(* IEC 61131-3 sources: 2026_Projet_YGO_ExcavatriceDragage/TOOLS/TEST_AUTO_CI/RESULTS/L_SIMULATION/tests (part 5) *)

(* ---- test_sim_manual_reference.st ---- *)
(* Copy-out explicite VAR_IN_OUT : le runner multi-FB sans source homonyme ne fait pas le post-traitement monobloc.
   Aucune valeur de reference inventee : seuls les resultats publics des FB sont restitues. *)
(* T418 : trois commandes IHM de reference, vrais codeurs/benne avec retours SimBench.
   Harnais des composants et routage explicite equivalent PRG, pas execution complete PLC.
   Aucun statut Homed/Reference positif n'est injecte. *)
SETUP
VAR
    bench : FB_SimBench;
    encoderM1 : FB_Encoder;
    encoderM2 : FB_Encoder;
    bucket : FB_Bucket;
    home : FB_CycleMachineHoming;
    cfgEncoder : ST_fbEncoder_Cfg;
    cfgBucket : ST_fbBucket_Config;
    calibM1 : ST_Encoder_Calib;
    calibM2 : ST_Encoder_Calib;
    hw1 : ST_fbEncoder_HwIn;
    hw2 : ST_fbEncoder_HwIn;
    bucketState : ST_fbBucket_State;
    bucketEdge : R_TRIG;
    raw1 : UDINT;
    raw2 : UDINT;
    btnM1 : BOOL;
    btnM2 : BOOL;
    btnBucket : BOOL;
END_VAR
END_SETUP

TEST 'TC-T418-REF-001 Trois commandes IHM etablissent les references dans le banc'
raw1 := 100000; raw2 := 200000; btnM1 := FALSE; btnM2 := FALSE; btnBucket := FALSE;
calibM1.Homed := FALSE; calibM2.Homed := FALSE; bucketState.BucketReferenced := FALSE;
cfgEncoder.PresetConfirmMode := E_PresetConfirmMode.READBACK_ONLY;
cfgBucket.OffsetOpenM := 2.25; cfgBucket.OffsetCloseM := 15.0; cfgBucket.CoherenceLimitM := 1.0;
bench.Enable := TRUE; home.Enable := TRUE; home.BootReady := TRUE; home.Mode := E_Mode.MAINT_N2; home.WinchesMechanicallyStopped := TRUE;
ADVANCE_TIME(10000000);
bench(M1_PresetTriggerCmd := encoderM1.HwOut.PresetTriggerCmd, M1_PresetValueOut := encoderM1.HwOut.PresetValueOut, M2_PresetTriggerCmd := encoderM2.HwOut.PresetTriggerCmd, M2_PresetValueOut := encoderM2.HwOut.PresetValueOut, RawPosM1 := raw1, RawPosM2 := raw2); raw1 := bench.RawPosM1; raw2 := bench.RawPosM2;
hw1.RawPosIn := bench.Winch.COD1_PosValue; hw1.SlaveOperational := TRUE; hw2.RawPosIn := bench.Winch.COD2_PosValue; hw2.SlaveOperational := TRUE;
encoderM1(Enable := TRUE, HomingPermit := TRUE, HomingAtTargetM := btnM1, CfgHomingTargetM := 8.7, CfgTopSensorPosM := 8.7, HwIn := hw1, Cfg := cfgEncoder, Calib := calibM1); calibM1 := encoderM1.Calib;
bucketEdge(CLK := btnBucket);
encoderM2(Enable := TRUE, HomingPermit := TRUE, HomingAtTargetM := btnM2 OR bucketEdge.Q, CfgHomingTargetM := 23.7, CfgTopSensorPosM := 23.7, UseDynamicTarget := bucketEdge.Q, DynamicHomingTargetM := encoderM1.Measurement.CablePosM + cfgBucket.OffsetCloseM, HwIn := hw2, Cfg := cfgEncoder, Calib := calibM2); calibM2 := encoderM2.Calib;
bucket(Enable := TRUE, Mode := E_Mode.MAINT_N2, PowerContactorEngaged := TRUE, CablePosM1 := encoderM1.Measurement.CablePosM, CablePosM2 := encoderM2.Measurement.CablePosM, HomedM1 := encoderM1.Homed, HomedM2 := encoderM2.Homed, HomedAndReliableM1 := encoderM1.HomedAndReliable, HomedAndReliableM2 := encoderM2.HomedAndReliable, HomingSuspectM1 := encoderM1.HomingSuspect, HomingSuspectM2 := encoderM2.HomingSuspect, ConfirmClosePosition := btnBucket, Config := cfgBucket, BucketState := bucketState); bucketState := bucket.BucketState;
home.M1Status.HomedAndReliable := encoderM1.HomedAndReliable; home.M2Status.HomedAndReliable := encoderM2.HomedAndReliable; home(BucketOffsetValid := bucketState.BucketReferenced, BtnValidation := bench.Operator.JoyBtnRaw);
ADVANCE_TIME(10000000);
bench(M1_PresetTriggerCmd := encoderM1.HwOut.PresetTriggerCmd, M1_PresetValueOut := encoderM1.HwOut.PresetValueOut, M2_PresetTriggerCmd := encoderM2.HwOut.PresetTriggerCmd, M2_PresetValueOut := encoderM2.HwOut.PresetValueOut, RawPosM1 := raw1, RawPosM2 := raw2); raw1 := bench.RawPosM1; raw2 := bench.RawPosM2;
hw1.RawPosIn := bench.Winch.COD1_PosValue; hw1.SlaveOperational := TRUE; hw2.RawPosIn := bench.Winch.COD2_PosValue; hw2.SlaveOperational := TRUE;
encoderM1(Enable := TRUE, HomingPermit := TRUE, HomingAtTargetM := btnM1, CfgHomingTargetM := 8.7, CfgTopSensorPosM := 8.7, HwIn := hw1, Cfg := cfgEncoder, Calib := calibM1); calibM1 := encoderM1.Calib;
bucketEdge(CLK := btnBucket);
encoderM2(Enable := TRUE, HomingPermit := TRUE, HomingAtTargetM := btnM2 OR bucketEdge.Q, CfgHomingTargetM := 23.7, CfgTopSensorPosM := 23.7, UseDynamicTarget := bucketEdge.Q, DynamicHomingTargetM := encoderM1.Measurement.CablePosM + cfgBucket.OffsetCloseM, HwIn := hw2, Cfg := cfgEncoder, Calib := calibM2); calibM2 := encoderM2.Calib;
bucket(Enable := TRUE, Mode := E_Mode.MAINT_N2, PowerContactorEngaged := TRUE, CablePosM1 := encoderM1.Measurement.CablePosM, CablePosM2 := encoderM2.Measurement.CablePosM, HomedM1 := encoderM1.Homed, HomedM2 := encoderM2.Homed, HomedAndReliableM1 := encoderM1.HomedAndReliable, HomedAndReliableM2 := encoderM2.HomedAndReliable, HomingSuspectM1 := encoderM1.HomingSuspect, HomingSuspectM2 := encoderM2.HomingSuspect, ConfirmClosePosition := btnBucket, Config := cfgBucket, BucketState := bucketState); bucketState := bucket.BucketState;
home.M1Status.HomedAndReliable := encoderM1.HomedAndReliable; home.M2Status.HomedAndReliable := encoderM2.HomedAndReliable; home(BucketOffsetValid := bucketState.BucketReferenced, BtnValidation := bench.Operator.JoyBtnRaw);
ASSERT_FALSE(home.MachineHomed, 'Boot non reference'); ASSERT_FALSE(encoderM1.Homed, 'M1 initial non reference'); ASSERT_FALSE(encoderM2.Homed, 'M2 initial non reference');
btnM1 := TRUE;
ADVANCE_TIME(10000000);
bench(M1_PresetTriggerCmd := encoderM1.HwOut.PresetTriggerCmd, M1_PresetValueOut := encoderM1.HwOut.PresetValueOut, M2_PresetTriggerCmd := encoderM2.HwOut.PresetTriggerCmd, M2_PresetValueOut := encoderM2.HwOut.PresetValueOut, RawPosM1 := raw1, RawPosM2 := raw2); raw1 := bench.RawPosM1; raw2 := bench.RawPosM2;
hw1.RawPosIn := bench.Winch.COD1_PosValue; hw1.SlaveOperational := TRUE; hw2.RawPosIn := bench.Winch.COD2_PosValue; hw2.SlaveOperational := TRUE;
encoderM1(Enable := TRUE, HomingPermit := TRUE, HomingAtTargetM := btnM1, CfgHomingTargetM := 8.7, CfgTopSensorPosM := 8.7, HwIn := hw1, Cfg := cfgEncoder, Calib := calibM1); calibM1 := encoderM1.Calib;
bucketEdge(CLK := btnBucket);
encoderM2(Enable := TRUE, HomingPermit := TRUE, HomingAtTargetM := btnM2 OR bucketEdge.Q, CfgHomingTargetM := 23.7, CfgTopSensorPosM := 23.7, UseDynamicTarget := bucketEdge.Q, DynamicHomingTargetM := encoderM1.Measurement.CablePosM + cfgBucket.OffsetCloseM, HwIn := hw2, Cfg := cfgEncoder, Calib := calibM2); calibM2 := encoderM2.Calib;
bucket(Enable := TRUE, Mode := E_Mode.MAINT_N2, PowerContactorEngaged := TRUE, CablePosM1 := encoderM1.Measurement.CablePosM, CablePosM2 := encoderM2.Measurement.CablePosM, HomedM1 := encoderM1.Homed, HomedM2 := encoderM2.Homed, HomedAndReliableM1 := encoderM1.HomedAndReliable, HomedAndReliableM2 := encoderM2.HomedAndReliable, HomingSuspectM1 := encoderM1.HomingSuspect, HomingSuspectM2 := encoderM2.HomingSuspect, ConfirmClosePosition := btnBucket, Config := cfgBucket, BucketState := bucketState); bucketState := bucket.BucketState;
home.M1Status.HomedAndReliable := encoderM1.HomedAndReliable; home.M2Status.HomedAndReliable := encoderM2.HomedAndReliable; home(BucketOffsetValid := bucketState.BucketReferenced, BtnValidation := bench.Operator.JoyBtnRaw);
btnM1 := FALSE;
ADVANCE_TIME(10000000);
bench(M1_PresetTriggerCmd := encoderM1.HwOut.PresetTriggerCmd, M1_PresetValueOut := encoderM1.HwOut.PresetValueOut, M2_PresetTriggerCmd := encoderM2.HwOut.PresetTriggerCmd, M2_PresetValueOut := encoderM2.HwOut.PresetValueOut, RawPosM1 := raw1, RawPosM2 := raw2); raw1 := bench.RawPosM1; raw2 := bench.RawPosM2;
hw1.RawPosIn := bench.Winch.COD1_PosValue; hw1.SlaveOperational := TRUE; hw2.RawPosIn := bench.Winch.COD2_PosValue; hw2.SlaveOperational := TRUE;
encoderM1(Enable := TRUE, HomingPermit := TRUE, HomingAtTargetM := btnM1, CfgHomingTargetM := 8.7, CfgTopSensorPosM := 8.7, HwIn := hw1, Cfg := cfgEncoder, Calib := calibM1); calibM1 := encoderM1.Calib;
bucketEdge(CLK := btnBucket);
encoderM2(Enable := TRUE, HomingPermit := TRUE, HomingAtTargetM := btnM2 OR bucketEdge.Q, CfgHomingTargetM := 23.7, CfgTopSensorPosM := 23.7, UseDynamicTarget := bucketEdge.Q, DynamicHomingTargetM := encoderM1.Measurement.CablePosM + cfgBucket.OffsetCloseM, HwIn := hw2, Cfg := cfgEncoder, Calib := calibM2); calibM2 := encoderM2.Calib;
bucket(Enable := TRUE, Mode := E_Mode.MAINT_N2, PowerContactorEngaged := TRUE, CablePosM1 := encoderM1.Measurement.CablePosM, CablePosM2 := encoderM2.Measurement.CablePosM, HomedM1 := encoderM1.Homed, HomedM2 := encoderM2.Homed, HomedAndReliableM1 := encoderM1.HomedAndReliable, HomedAndReliableM2 := encoderM2.HomedAndReliable, HomingSuspectM1 := encoderM1.HomingSuspect, HomingSuspectM2 := encoderM2.HomingSuspect, ConfirmClosePosition := btnBucket, Config := cfgBucket, BucketState := bucketState); bucketState := bucket.BucketState;
home.M1Status.HomedAndReliable := encoderM1.HomedAndReliable; home.M2Status.HomedAndReliable := encoderM2.HomedAndReliable; home(BucketOffsetValid := bucketState.BucketReferenced, BtnValidation := bench.Operator.JoyBtnRaw);
ADVANCE_TIME(10000000);
bench(M1_PresetTriggerCmd := encoderM1.HwOut.PresetTriggerCmd, M1_PresetValueOut := encoderM1.HwOut.PresetValueOut, M2_PresetTriggerCmd := encoderM2.HwOut.PresetTriggerCmd, M2_PresetValueOut := encoderM2.HwOut.PresetValueOut, RawPosM1 := raw1, RawPosM2 := raw2); raw1 := bench.RawPosM1; raw2 := bench.RawPosM2;
hw1.RawPosIn := bench.Winch.COD1_PosValue; hw1.SlaveOperational := TRUE; hw2.RawPosIn := bench.Winch.COD2_PosValue; hw2.SlaveOperational := TRUE;
encoderM1(Enable := TRUE, HomingPermit := TRUE, HomingAtTargetM := btnM1, CfgHomingTargetM := 8.7, CfgTopSensorPosM := 8.7, HwIn := hw1, Cfg := cfgEncoder, Calib := calibM1); calibM1 := encoderM1.Calib;
bucketEdge(CLK := btnBucket);
encoderM2(Enable := TRUE, HomingPermit := TRUE, HomingAtTargetM := btnM2 OR bucketEdge.Q, CfgHomingTargetM := 23.7, CfgTopSensorPosM := 23.7, UseDynamicTarget := bucketEdge.Q, DynamicHomingTargetM := encoderM1.Measurement.CablePosM + cfgBucket.OffsetCloseM, HwIn := hw2, Cfg := cfgEncoder, Calib := calibM2); calibM2 := encoderM2.Calib;
bucket(Enable := TRUE, Mode := E_Mode.MAINT_N2, PowerContactorEngaged := TRUE, CablePosM1 := encoderM1.Measurement.CablePosM, CablePosM2 := encoderM2.Measurement.CablePosM, HomedM1 := encoderM1.Homed, HomedM2 := encoderM2.Homed, HomedAndReliableM1 := encoderM1.HomedAndReliable, HomedAndReliableM2 := encoderM2.HomedAndReliable, HomingSuspectM1 := encoderM1.HomingSuspect, HomingSuspectM2 := encoderM2.HomingSuspect, ConfirmClosePosition := btnBucket, Config := cfgBucket, BucketState := bucketState); bucketState := bucket.BucketState;
home.M1Status.HomedAndReliable := encoderM1.HomedAndReliable; home.M2Status.HomedAndReliable := encoderM2.HomedAndReliable; home(BucketOffsetValid := bucketState.BucketReferenced, BtnValidation := bench.Operator.JoyBtnRaw);
ADVANCE_TIME(10000000);
bench(M1_PresetTriggerCmd := encoderM1.HwOut.PresetTriggerCmd, M1_PresetValueOut := encoderM1.HwOut.PresetValueOut, M2_PresetTriggerCmd := encoderM2.HwOut.PresetTriggerCmd, M2_PresetValueOut := encoderM2.HwOut.PresetValueOut, RawPosM1 := raw1, RawPosM2 := raw2); raw1 := bench.RawPosM1; raw2 := bench.RawPosM2;
hw1.RawPosIn := bench.Winch.COD1_PosValue; hw1.SlaveOperational := TRUE; hw2.RawPosIn := bench.Winch.COD2_PosValue; hw2.SlaveOperational := TRUE;
encoderM1(Enable := TRUE, HomingPermit := TRUE, HomingAtTargetM := btnM1, CfgHomingTargetM := 8.7, CfgTopSensorPosM := 8.7, HwIn := hw1, Cfg := cfgEncoder, Calib := calibM1); calibM1 := encoderM1.Calib;
bucketEdge(CLK := btnBucket);
encoderM2(Enable := TRUE, HomingPermit := TRUE, HomingAtTargetM := btnM2 OR bucketEdge.Q, CfgHomingTargetM := 23.7, CfgTopSensorPosM := 23.7, UseDynamicTarget := bucketEdge.Q, DynamicHomingTargetM := encoderM1.Measurement.CablePosM + cfgBucket.OffsetCloseM, HwIn := hw2, Cfg := cfgEncoder, Calib := calibM2); calibM2 := encoderM2.Calib;
bucket(Enable := TRUE, Mode := E_Mode.MAINT_N2, PowerContactorEngaged := TRUE, CablePosM1 := encoderM1.Measurement.CablePosM, CablePosM2 := encoderM2.Measurement.CablePosM, HomedM1 := encoderM1.Homed, HomedM2 := encoderM2.Homed, HomedAndReliableM1 := encoderM1.HomedAndReliable, HomedAndReliableM2 := encoderM2.HomedAndReliable, HomingSuspectM1 := encoderM1.HomingSuspect, HomingSuspectM2 := encoderM2.HomingSuspect, ConfirmClosePosition := btnBucket, Config := cfgBucket, BucketState := bucketState); bucketState := bucket.BucketState;
home.M1Status.HomedAndReliable := encoderM1.HomedAndReliable; home.M2Status.HomedAndReliable := encoderM2.HomedAndReliable; home(BucketOffsetValid := bucketState.BucketReferenced, BtnValidation := bench.Operator.JoyBtnRaw);
ADVANCE_TIME(10000000);
bench(M1_PresetTriggerCmd := encoderM1.HwOut.PresetTriggerCmd, M1_PresetValueOut := encoderM1.HwOut.PresetValueOut, M2_PresetTriggerCmd := encoderM2.HwOut.PresetTriggerCmd, M2_PresetValueOut := encoderM2.HwOut.PresetValueOut, RawPosM1 := raw1, RawPosM2 := raw2); raw1 := bench.RawPosM1; raw2 := bench.RawPosM2;
hw1.RawPosIn := bench.Winch.COD1_PosValue; hw1.SlaveOperational := TRUE; hw2.RawPosIn := bench.Winch.COD2_PosValue; hw2.SlaveOperational := TRUE;
encoderM1(Enable := TRUE, HomingPermit := TRUE, HomingAtTargetM := btnM1, CfgHomingTargetM := 8.7, CfgTopSensorPosM := 8.7, HwIn := hw1, Cfg := cfgEncoder, Calib := calibM1); calibM1 := encoderM1.Calib;
bucketEdge(CLK := btnBucket);
encoderM2(Enable := TRUE, HomingPermit := TRUE, HomingAtTargetM := btnM2 OR bucketEdge.Q, CfgHomingTargetM := 23.7, CfgTopSensorPosM := 23.7, UseDynamicTarget := bucketEdge.Q, DynamicHomingTargetM := encoderM1.Measurement.CablePosM + cfgBucket.OffsetCloseM, HwIn := hw2, Cfg := cfgEncoder, Calib := calibM2); calibM2 := encoderM2.Calib;
bucket(Enable := TRUE, Mode := E_Mode.MAINT_N2, PowerContactorEngaged := TRUE, CablePosM1 := encoderM1.Measurement.CablePosM, CablePosM2 := encoderM2.Measurement.CablePosM, HomedM1 := encoderM1.Homed, HomedM2 := encoderM2.Homed, HomedAndReliableM1 := encoderM1.HomedAndReliable, HomedAndReliableM2 := encoderM2.HomedAndReliable, HomingSuspectM1 := encoderM1.HomingSuspect, HomingSuspectM2 := encoderM2.HomingSuspect, ConfirmClosePosition := btnBucket, Config := cfgBucket, BucketState := bucketState); bucketState := bucket.BucketState;
home.M1Status.HomedAndReliable := encoderM1.HomedAndReliable; home.M2Status.HomedAndReliable := encoderM2.HomedAndReliable; home(BucketOffsetValid := bucketState.BucketReferenced, BtnValidation := bench.Operator.JoyBtnRaw);
ADVANCE_TIME(10000000);
bench(M1_PresetTriggerCmd := encoderM1.HwOut.PresetTriggerCmd, M1_PresetValueOut := encoderM1.HwOut.PresetValueOut, M2_PresetTriggerCmd := encoderM2.HwOut.PresetTriggerCmd, M2_PresetValueOut := encoderM2.HwOut.PresetValueOut, RawPosM1 := raw1, RawPosM2 := raw2); raw1 := bench.RawPosM1; raw2 := bench.RawPosM2;
hw1.RawPosIn := bench.Winch.COD1_PosValue; hw1.SlaveOperational := TRUE; hw2.RawPosIn := bench.Winch.COD2_PosValue; hw2.SlaveOperational := TRUE;
encoderM1(Enable := TRUE, HomingPermit := TRUE, HomingAtTargetM := btnM1, CfgHomingTargetM := 8.7, CfgTopSensorPosM := 8.7, HwIn := hw1, Cfg := cfgEncoder, Calib := calibM1); calibM1 := encoderM1.Calib;
bucketEdge(CLK := btnBucket);
encoderM2(Enable := TRUE, HomingPermit := TRUE, HomingAtTargetM := btnM2 OR bucketEdge.Q, CfgHomingTargetM := 23.7, CfgTopSensorPosM := 23.7, UseDynamicTarget := bucketEdge.Q, DynamicHomingTargetM := encoderM1.Measurement.CablePosM + cfgBucket.OffsetCloseM, HwIn := hw2, Cfg := cfgEncoder, Calib := calibM2); calibM2 := encoderM2.Calib;
bucket(Enable := TRUE, Mode := E_Mode.MAINT_N2, PowerContactorEngaged := TRUE, CablePosM1 := encoderM1.Measurement.CablePosM, CablePosM2 := encoderM2.Measurement.CablePosM, HomedM1 := encoderM1.Homed, HomedM2 := encoderM2.Homed, HomedAndReliableM1 := encoderM1.HomedAndReliable, HomedAndReliableM2 := encoderM2.HomedAndReliable, HomingSuspectM1 := encoderM1.HomingSuspect, HomingSuspectM2 := encoderM2.HomingSuspect, ConfirmClosePosition := btnBucket, Config := cfgBucket, BucketState := bucketState); bucketState := bucket.BucketState;
home.M1Status.HomedAndReliable := encoderM1.HomedAndReliable; home.M2Status.HomedAndReliable := encoderM2.HomedAndReliable; home(BucketOffsetValid := bucketState.BucketReferenced, BtnValidation := bench.Operator.JoyBtnRaw);
ADVANCE_TIME(10000000);
bench(M1_PresetTriggerCmd := encoderM1.HwOut.PresetTriggerCmd, M1_PresetValueOut := encoderM1.HwOut.PresetValueOut, M2_PresetTriggerCmd := encoderM2.HwOut.PresetTriggerCmd, M2_PresetValueOut := encoderM2.HwOut.PresetValueOut, RawPosM1 := raw1, RawPosM2 := raw2); raw1 := bench.RawPosM1; raw2 := bench.RawPosM2;
hw1.RawPosIn := bench.Winch.COD1_PosValue; hw1.SlaveOperational := TRUE; hw2.RawPosIn := bench.Winch.COD2_PosValue; hw2.SlaveOperational := TRUE;
encoderM1(Enable := TRUE, HomingPermit := TRUE, HomingAtTargetM := btnM1, CfgHomingTargetM := 8.7, CfgTopSensorPosM := 8.7, HwIn := hw1, Cfg := cfgEncoder, Calib := calibM1); calibM1 := encoderM1.Calib;
bucketEdge(CLK := btnBucket);
encoderM2(Enable := TRUE, HomingPermit := TRUE, HomingAtTargetM := btnM2 OR bucketEdge.Q, CfgHomingTargetM := 23.7, CfgTopSensorPosM := 23.7, UseDynamicTarget := bucketEdge.Q, DynamicHomingTargetM := encoderM1.Measurement.CablePosM + cfgBucket.OffsetCloseM, HwIn := hw2, Cfg := cfgEncoder, Calib := calibM2); calibM2 := encoderM2.Calib;
bucket(Enable := TRUE, Mode := E_Mode.MAINT_N2, PowerContactorEngaged := TRUE, CablePosM1 := encoderM1.Measurement.CablePosM, CablePosM2 := encoderM2.Measurement.CablePosM, HomedM1 := encoderM1.Homed, HomedM2 := encoderM2.Homed, HomedAndReliableM1 := encoderM1.HomedAndReliable, HomedAndReliableM2 := encoderM2.HomedAndReliable, HomingSuspectM1 := encoderM1.HomingSuspect, HomingSuspectM2 := encoderM2.HomingSuspect, ConfirmClosePosition := btnBucket, Config := cfgBucket, BucketState := bucketState); bucketState := bucket.BucketState;
home.M1Status.HomedAndReliable := encoderM1.HomedAndReliable; home.M2Status.HomedAndReliable := encoderM2.HomedAndReliable; home(BucketOffsetValid := bucketState.BucketReferenced, BtnValidation := bench.Operator.JoyBtnRaw);
ADVANCE_TIME(10000000);
bench(M1_PresetTriggerCmd := encoderM1.HwOut.PresetTriggerCmd, M1_PresetValueOut := encoderM1.HwOut.PresetValueOut, M2_PresetTriggerCmd := encoderM2.HwOut.PresetTriggerCmd, M2_PresetValueOut := encoderM2.HwOut.PresetValueOut, RawPosM1 := raw1, RawPosM2 := raw2); raw1 := bench.RawPosM1; raw2 := bench.RawPosM2;
hw1.RawPosIn := bench.Winch.COD1_PosValue; hw1.SlaveOperational := TRUE; hw2.RawPosIn := bench.Winch.COD2_PosValue; hw2.SlaveOperational := TRUE;
encoderM1(Enable := TRUE, HomingPermit := TRUE, HomingAtTargetM := btnM1, CfgHomingTargetM := 8.7, CfgTopSensorPosM := 8.7, HwIn := hw1, Cfg := cfgEncoder, Calib := calibM1); calibM1 := encoderM1.Calib;
bucketEdge(CLK := btnBucket);
encoderM2(Enable := TRUE, HomingPermit := TRUE, HomingAtTargetM := btnM2 OR bucketEdge.Q, CfgHomingTargetM := 23.7, CfgTopSensorPosM := 23.7, UseDynamicTarget := bucketEdge.Q, DynamicHomingTargetM := encoderM1.Measurement.CablePosM + cfgBucket.OffsetCloseM, HwIn := hw2, Cfg := cfgEncoder, Calib := calibM2); calibM2 := encoderM2.Calib;
bucket(Enable := TRUE, Mode := E_Mode.MAINT_N2, PowerContactorEngaged := TRUE, CablePosM1 := encoderM1.Measurement.CablePosM, CablePosM2 := encoderM2.Measurement.CablePosM, HomedM1 := encoderM1.Homed, HomedM2 := encoderM2.Homed, HomedAndReliableM1 := encoderM1.HomedAndReliable, HomedAndReliableM2 := encoderM2.HomedAndReliable, HomingSuspectM1 := encoderM1.HomingSuspect, HomingSuspectM2 := encoderM2.HomingSuspect, ConfirmClosePosition := btnBucket, Config := cfgBucket, BucketState := bucketState); bucketState := bucket.BucketState;
home.M1Status.HomedAndReliable := encoderM1.HomedAndReliable; home.M2Status.HomedAndReliable := encoderM2.HomedAndReliable; home(BucketOffsetValid := bucketState.BucketReferenced, BtnValidation := bench.Operator.JoyBtnRaw);
ADVANCE_TIME(10000000);
bench(M1_PresetTriggerCmd := encoderM1.HwOut.PresetTriggerCmd, M1_PresetValueOut := encoderM1.HwOut.PresetValueOut, M2_PresetTriggerCmd := encoderM2.HwOut.PresetTriggerCmd, M2_PresetValueOut := encoderM2.HwOut.PresetValueOut, RawPosM1 := raw1, RawPosM2 := raw2); raw1 := bench.RawPosM1; raw2 := bench.RawPosM2;
hw1.RawPosIn := bench.Winch.COD1_PosValue; hw1.SlaveOperational := TRUE; hw2.RawPosIn := bench.Winch.COD2_PosValue; hw2.SlaveOperational := TRUE;
encoderM1(Enable := TRUE, HomingPermit := TRUE, HomingAtTargetM := btnM1, CfgHomingTargetM := 8.7, CfgTopSensorPosM := 8.7, HwIn := hw1, Cfg := cfgEncoder, Calib := calibM1); calibM1 := encoderM1.Calib;
bucketEdge(CLK := btnBucket);
encoderM2(Enable := TRUE, HomingPermit := TRUE, HomingAtTargetM := btnM2 OR bucketEdge.Q, CfgHomingTargetM := 23.7, CfgTopSensorPosM := 23.7, UseDynamicTarget := bucketEdge.Q, DynamicHomingTargetM := encoderM1.Measurement.CablePosM + cfgBucket.OffsetCloseM, HwIn := hw2, Cfg := cfgEncoder, Calib := calibM2); calibM2 := encoderM2.Calib;
bucket(Enable := TRUE, Mode := E_Mode.MAINT_N2, PowerContactorEngaged := TRUE, CablePosM1 := encoderM1.Measurement.CablePosM, CablePosM2 := encoderM2.Measurement.CablePosM, HomedM1 := encoderM1.Homed, HomedM2 := encoderM2.Homed, HomedAndReliableM1 := encoderM1.HomedAndReliable, HomedAndReliableM2 := encoderM2.HomedAndReliable, HomingSuspectM1 := encoderM1.HomingSuspect, HomingSuspectM2 := encoderM2.HomingSuspect, ConfirmClosePosition := btnBucket, Config := cfgBucket, BucketState := bucketState); bucketState := bucket.BucketState;
home.M1Status.HomedAndReliable := encoderM1.HomedAndReliable; home.M2Status.HomedAndReliable := encoderM2.HomedAndReliable; home(BucketOffsetValid := bucketState.BucketReferenced, BtnValidation := bench.Operator.JoyBtnRaw);
ADVANCE_TIME(10000000);
bench(M1_PresetTriggerCmd := encoderM1.HwOut.PresetTriggerCmd, M1_PresetValueOut := encoderM1.HwOut.PresetValueOut, M2_PresetTriggerCmd := encoderM2.HwOut.PresetTriggerCmd, M2_PresetValueOut := encoderM2.HwOut.PresetValueOut, RawPosM1 := raw1, RawPosM2 := raw2); raw1 := bench.RawPosM1; raw2 := bench.RawPosM2;
hw1.RawPosIn := bench.Winch.COD1_PosValue; hw1.SlaveOperational := TRUE; hw2.RawPosIn := bench.Winch.COD2_PosValue; hw2.SlaveOperational := TRUE;
encoderM1(Enable := TRUE, HomingPermit := TRUE, HomingAtTargetM := btnM1, CfgHomingTargetM := 8.7, CfgTopSensorPosM := 8.7, HwIn := hw1, Cfg := cfgEncoder, Calib := calibM1); calibM1 := encoderM1.Calib;
bucketEdge(CLK := btnBucket);
encoderM2(Enable := TRUE, HomingPermit := TRUE, HomingAtTargetM := btnM2 OR bucketEdge.Q, CfgHomingTargetM := 23.7, CfgTopSensorPosM := 23.7, UseDynamicTarget := bucketEdge.Q, DynamicHomingTargetM := encoderM1.Measurement.CablePosM + cfgBucket.OffsetCloseM, HwIn := hw2, Cfg := cfgEncoder, Calib := calibM2); calibM2 := encoderM2.Calib;
bucket(Enable := TRUE, Mode := E_Mode.MAINT_N2, PowerContactorEngaged := TRUE, CablePosM1 := encoderM1.Measurement.CablePosM, CablePosM2 := encoderM2.Measurement.CablePosM, HomedM1 := encoderM1.Homed, HomedM2 := encoderM2.Homed, HomedAndReliableM1 := encoderM1.HomedAndReliable, HomedAndReliableM2 := encoderM2.HomedAndReliable, HomingSuspectM1 := encoderM1.HomingSuspect, HomingSuspectM2 := encoderM2.HomingSuspect, ConfirmClosePosition := btnBucket, Config := cfgBucket, BucketState := bucketState); bucketState := bucket.BucketState;
home.M1Status.HomedAndReliable := encoderM1.HomedAndReliable; home.M2Status.HomedAndReliable := encoderM2.HomedAndReliable; home(BucketOffsetValid := bucketState.BucketReferenced, BtnValidation := bench.Operator.JoyBtnRaw);
ADVANCE_TIME(10000000);
bench(M1_PresetTriggerCmd := encoderM1.HwOut.PresetTriggerCmd, M1_PresetValueOut := encoderM1.HwOut.PresetValueOut, M2_PresetTriggerCmd := encoderM2.HwOut.PresetTriggerCmd, M2_PresetValueOut := encoderM2.HwOut.PresetValueOut, RawPosM1 := raw1, RawPosM2 := raw2); raw1 := bench.RawPosM1; raw2 := bench.RawPosM2;
hw1.RawPosIn := bench.Winch.COD1_PosValue; hw1.SlaveOperational := TRUE; hw2.RawPosIn := bench.Winch.COD2_PosValue; hw2.SlaveOperational := TRUE;
encoderM1(Enable := TRUE, HomingPermit := TRUE, HomingAtTargetM := btnM1, CfgHomingTargetM := 8.7, CfgTopSensorPosM := 8.7, HwIn := hw1, Cfg := cfgEncoder, Calib := calibM1); calibM1 := encoderM1.Calib;
bucketEdge(CLK := btnBucket);
encoderM2(Enable := TRUE, HomingPermit := TRUE, HomingAtTargetM := btnM2 OR bucketEdge.Q, CfgHomingTargetM := 23.7, CfgTopSensorPosM := 23.7, UseDynamicTarget := bucketEdge.Q, DynamicHomingTargetM := encoderM1.Measurement.CablePosM + cfgBucket.OffsetCloseM, HwIn := hw2, Cfg := cfgEncoder, Calib := calibM2); calibM2 := encoderM2.Calib;
bucket(Enable := TRUE, Mode := E_Mode.MAINT_N2, PowerContactorEngaged := TRUE, CablePosM1 := encoderM1.Measurement.CablePosM, CablePosM2 := encoderM2.Measurement.CablePosM, HomedM1 := encoderM1.Homed, HomedM2 := encoderM2.Homed, HomedAndReliableM1 := encoderM1.HomedAndReliable, HomedAndReliableM2 := encoderM2.HomedAndReliable, HomingSuspectM1 := encoderM1.HomingSuspect, HomingSuspectM2 := encoderM2.HomingSuspect, ConfirmClosePosition := btnBucket, Config := cfgBucket, BucketState := bucketState); bucketState := bucket.BucketState;
home.M1Status.HomedAndReliable := encoderM1.HomedAndReliable; home.M2Status.HomedAndReliable := encoderM2.HomedAndReliable; home(BucketOffsetValid := bucketState.BucketReferenced, BtnValidation := bench.Operator.JoyBtnRaw);
ADVANCE_TIME(10000000);
bench(M1_PresetTriggerCmd := encoderM1.HwOut.PresetTriggerCmd, M1_PresetValueOut := encoderM1.HwOut.PresetValueOut, M2_PresetTriggerCmd := encoderM2.HwOut.PresetTriggerCmd, M2_PresetValueOut := encoderM2.HwOut.PresetValueOut, RawPosM1 := raw1, RawPosM2 := raw2); raw1 := bench.RawPosM1; raw2 := bench.RawPosM2;
hw1.RawPosIn := bench.Winch.COD1_PosValue; hw1.SlaveOperational := TRUE; hw2.RawPosIn := bench.Winch.COD2_PosValue; hw2.SlaveOperational := TRUE;
encoderM1(Enable := TRUE, HomingPermit := TRUE, HomingAtTargetM := btnM1, CfgHomingTargetM := 8.7, CfgTopSensorPosM := 8.7, HwIn := hw1, Cfg := cfgEncoder, Calib := calibM1); calibM1 := encoderM1.Calib;
bucketEdge(CLK := btnBucket);
encoderM2(Enable := TRUE, HomingPermit := TRUE, HomingAtTargetM := btnM2 OR bucketEdge.Q, CfgHomingTargetM := 23.7, CfgTopSensorPosM := 23.7, UseDynamicTarget := bucketEdge.Q, DynamicHomingTargetM := encoderM1.Measurement.CablePosM + cfgBucket.OffsetCloseM, HwIn := hw2, Cfg := cfgEncoder, Calib := calibM2); calibM2 := encoderM2.Calib;
bucket(Enable := TRUE, Mode := E_Mode.MAINT_N2, PowerContactorEngaged := TRUE, CablePosM1 := encoderM1.Measurement.CablePosM, CablePosM2 := encoderM2.Measurement.CablePosM, HomedM1 := encoderM1.Homed, HomedM2 := encoderM2.Homed, HomedAndReliableM1 := encoderM1.HomedAndReliable, HomedAndReliableM2 := encoderM2.HomedAndReliable, HomingSuspectM1 := encoderM1.HomingSuspect, HomingSuspectM2 := encoderM2.HomingSuspect, ConfirmClosePosition := btnBucket, Config := cfgBucket, BucketState := bucketState); bucketState := bucket.BucketState;
home.M1Status.HomedAndReliable := encoderM1.HomedAndReliable; home.M2Status.HomedAndReliable := encoderM2.HomedAndReliable; home(BucketOffsetValid := bucketState.BucketReferenced, BtnValidation := bench.Operator.JoyBtnRaw);
ADVANCE_TIME(10000000);
bench(M1_PresetTriggerCmd := encoderM1.HwOut.PresetTriggerCmd, M1_PresetValueOut := encoderM1.HwOut.PresetValueOut, M2_PresetTriggerCmd := encoderM2.HwOut.PresetTriggerCmd, M2_PresetValueOut := encoderM2.HwOut.PresetValueOut, RawPosM1 := raw1, RawPosM2 := raw2); raw1 := bench.RawPosM1; raw2 := bench.RawPosM2;
hw1.RawPosIn := bench.Winch.COD1_PosValue; hw1.SlaveOperational := TRUE; hw2.RawPosIn := bench.Winch.COD2_PosValue; hw2.SlaveOperational := TRUE;
encoderM1(Enable := TRUE, HomingPermit := TRUE, HomingAtTargetM := btnM1, CfgHomingTargetM := 8.7, CfgTopSensorPosM := 8.7, HwIn := hw1, Cfg := cfgEncoder, Calib := calibM1); calibM1 := encoderM1.Calib;
bucketEdge(CLK := btnBucket);
encoderM2(Enable := TRUE, HomingPermit := TRUE, HomingAtTargetM := btnM2 OR bucketEdge.Q, CfgHomingTargetM := 23.7, CfgTopSensorPosM := 23.7, UseDynamicTarget := bucketEdge.Q, DynamicHomingTargetM := encoderM1.Measurement.CablePosM + cfgBucket.OffsetCloseM, HwIn := hw2, Cfg := cfgEncoder, Calib := calibM2); calibM2 := encoderM2.Calib;
bucket(Enable := TRUE, Mode := E_Mode.MAINT_N2, PowerContactorEngaged := TRUE, CablePosM1 := encoderM1.Measurement.CablePosM, CablePosM2 := encoderM2.Measurement.CablePosM, HomedM1 := encoderM1.Homed, HomedM2 := encoderM2.Homed, HomedAndReliableM1 := encoderM1.HomedAndReliable, HomedAndReliableM2 := encoderM2.HomedAndReliable, HomingSuspectM1 := encoderM1.HomingSuspect, HomingSuspectM2 := encoderM2.HomingSuspect, ConfirmClosePosition := btnBucket, Config := cfgBucket, BucketState := bucketState); bucketState := bucket.BucketState;
home.M1Status.HomedAndReliable := encoderM1.HomedAndReliable; home.M2Status.HomedAndReliable := encoderM2.HomedAndReliable; home(BucketOffsetValid := bucketState.BucketReferenced, BtnValidation := bench.Operator.JoyBtnRaw);
ADVANCE_TIME(10000000);
bench(M1_PresetTriggerCmd := encoderM1.HwOut.PresetTriggerCmd, M1_PresetValueOut := encoderM1.HwOut.PresetValueOut, M2_PresetTriggerCmd := encoderM2.HwOut.PresetTriggerCmd, M2_PresetValueOut := encoderM2.HwOut.PresetValueOut, RawPosM1 := raw1, RawPosM2 := raw2); raw1 := bench.RawPosM1; raw2 := bench.RawPosM2;
hw1.RawPosIn := bench.Winch.COD1_PosValue; hw1.SlaveOperational := TRUE; hw2.RawPosIn := bench.Winch.COD2_PosValue; hw2.SlaveOperational := TRUE;
encoderM1(Enable := TRUE, HomingPermit := TRUE, HomingAtTargetM := btnM1, CfgHomingTargetM := 8.7, CfgTopSensorPosM := 8.7, HwIn := hw1, Cfg := cfgEncoder, Calib := calibM1); calibM1 := encoderM1.Calib;
bucketEdge(CLK := btnBucket);
encoderM2(Enable := TRUE, HomingPermit := TRUE, HomingAtTargetM := btnM2 OR bucketEdge.Q, CfgHomingTargetM := 23.7, CfgTopSensorPosM := 23.7, UseDynamicTarget := bucketEdge.Q, DynamicHomingTargetM := encoderM1.Measurement.CablePosM + cfgBucket.OffsetCloseM, HwIn := hw2, Cfg := cfgEncoder, Calib := calibM2); calibM2 := encoderM2.Calib;
bucket(Enable := TRUE, Mode := E_Mode.MAINT_N2, PowerContactorEngaged := TRUE, CablePosM1 := encoderM1.Measurement.CablePosM, CablePosM2 := encoderM2.Measurement.CablePosM, HomedM1 := encoderM1.Homed, HomedM2 := encoderM2.Homed, HomedAndReliableM1 := encoderM1.HomedAndReliable, HomedAndReliableM2 := encoderM2.HomedAndReliable, HomingSuspectM1 := encoderM1.HomingSuspect, HomingSuspectM2 := encoderM2.HomingSuspect, ConfirmClosePosition := btnBucket, Config := cfgBucket, BucketState := bucketState); bucketState := bucket.BucketState;
home.M1Status.HomedAndReliable := encoderM1.HomedAndReliable; home.M2Status.HomedAndReliable := encoderM2.HomedAndReliable; home(BucketOffsetValid := bucketState.BucketReferenced, BtnValidation := bench.Operator.JoyBtnRaw);
ADVANCE_TIME(10000000);
bench(M1_PresetTriggerCmd := encoderM1.HwOut.PresetTriggerCmd, M1_PresetValueOut := encoderM1.HwOut.PresetValueOut, M2_PresetTriggerCmd := encoderM2.HwOut.PresetTriggerCmd, M2_PresetValueOut := encoderM2.HwOut.PresetValueOut, RawPosM1 := raw1, RawPosM2 := raw2); raw1 := bench.RawPosM1; raw2 := bench.RawPosM2;
hw1.RawPosIn := bench.Winch.COD1_PosValue; hw1.SlaveOperational := TRUE; hw2.RawPosIn := bench.Winch.COD2_PosValue; hw2.SlaveOperational := TRUE;
encoderM1(Enable := TRUE, HomingPermit := TRUE, HomingAtTargetM := btnM1, CfgHomingTargetM := 8.7, CfgTopSensorPosM := 8.7, HwIn := hw1, Cfg := cfgEncoder, Calib := calibM1); calibM1 := encoderM1.Calib;
bucketEdge(CLK := btnBucket);
encoderM2(Enable := TRUE, HomingPermit := TRUE, HomingAtTargetM := btnM2 OR bucketEdge.Q, CfgHomingTargetM := 23.7, CfgTopSensorPosM := 23.7, UseDynamicTarget := bucketEdge.Q, DynamicHomingTargetM := encoderM1.Measurement.CablePosM + cfgBucket.OffsetCloseM, HwIn := hw2, Cfg := cfgEncoder, Calib := calibM2); calibM2 := encoderM2.Calib;
bucket(Enable := TRUE, Mode := E_Mode.MAINT_N2, PowerContactorEngaged := TRUE, CablePosM1 := encoderM1.Measurement.CablePosM, CablePosM2 := encoderM2.Measurement.CablePosM, HomedM1 := encoderM1.Homed, HomedM2 := encoderM2.Homed, HomedAndReliableM1 := encoderM1.HomedAndReliable, HomedAndReliableM2 := encoderM2.HomedAndReliable, HomingSuspectM1 := encoderM1.HomingSuspect, HomingSuspectM2 := encoderM2.HomingSuspect, ConfirmClosePosition := btnBucket, Config := cfgBucket, BucketState := bucketState); bucketState := bucket.BucketState;
home.M1Status.HomedAndReliable := encoderM1.HomedAndReliable; home.M2Status.HomedAndReliable := encoderM2.HomedAndReliable; home(BucketOffsetValid := bucketState.BucketReferenced, BtnValidation := bench.Operator.JoyBtnRaw);
ADVANCE_TIME(10000000);
bench(M1_PresetTriggerCmd := encoderM1.HwOut.PresetTriggerCmd, M1_PresetValueOut := encoderM1.HwOut.PresetValueOut, M2_PresetTriggerCmd := encoderM2.HwOut.PresetTriggerCmd, M2_PresetValueOut := encoderM2.HwOut.PresetValueOut, RawPosM1 := raw1, RawPosM2 := raw2); raw1 := bench.RawPosM1; raw2 := bench.RawPosM2;
hw1.RawPosIn := bench.Winch.COD1_PosValue; hw1.SlaveOperational := TRUE; hw2.RawPosIn := bench.Winch.COD2_PosValue; hw2.SlaveOperational := TRUE;
encoderM1(Enable := TRUE, HomingPermit := TRUE, HomingAtTargetM := btnM1, CfgHomingTargetM := 8.7, CfgTopSensorPosM := 8.7, HwIn := hw1, Cfg := cfgEncoder, Calib := calibM1); calibM1 := encoderM1.Calib;
bucketEdge(CLK := btnBucket);
encoderM2(Enable := TRUE, HomingPermit := TRUE, HomingAtTargetM := btnM2 OR bucketEdge.Q, CfgHomingTargetM := 23.7, CfgTopSensorPosM := 23.7, UseDynamicTarget := bucketEdge.Q, DynamicHomingTargetM := encoderM1.Measurement.CablePosM + cfgBucket.OffsetCloseM, HwIn := hw2, Cfg := cfgEncoder, Calib := calibM2); calibM2 := encoderM2.Calib;
bucket(Enable := TRUE, Mode := E_Mode.MAINT_N2, PowerContactorEngaged := TRUE, CablePosM1 := encoderM1.Measurement.CablePosM, CablePosM2 := encoderM2.Measurement.CablePosM, HomedM1 := encoderM1.Homed, HomedM2 := encoderM2.Homed, HomedAndReliableM1 := encoderM1.HomedAndReliable, HomedAndReliableM2 := encoderM2.HomedAndReliable, HomingSuspectM1 := encoderM1.HomingSuspect, HomingSuspectM2 := encoderM2.HomingSuspect, ConfirmClosePosition := btnBucket, Config := cfgBucket, BucketState := bucketState); bucketState := bucket.BucketState;
home.M1Status.HomedAndReliable := encoderM1.HomedAndReliable; home.M2Status.HomedAndReliable := encoderM2.HomedAndReliable; home(BucketOffsetValid := bucketState.BucketReferenced, BtnValidation := bench.Operator.JoyBtnRaw);
ADVANCE_TIME(10000000);
bench(M1_PresetTriggerCmd := encoderM1.HwOut.PresetTriggerCmd, M1_PresetValueOut := encoderM1.HwOut.PresetValueOut, M2_PresetTriggerCmd := encoderM2.HwOut.PresetTriggerCmd, M2_PresetValueOut := encoderM2.HwOut.PresetValueOut, RawPosM1 := raw1, RawPosM2 := raw2); raw1 := bench.RawPosM1; raw2 := bench.RawPosM2;
hw1.RawPosIn := bench.Winch.COD1_PosValue; hw1.SlaveOperational := TRUE; hw2.RawPosIn := bench.Winch.COD2_PosValue; hw2.SlaveOperational := TRUE;
encoderM1(Enable := TRUE, HomingPermit := TRUE, HomingAtTargetM := btnM1, CfgHomingTargetM := 8.7, CfgTopSensorPosM := 8.7, HwIn := hw1, Cfg := cfgEncoder, Calib := calibM1); calibM1 := encoderM1.Calib;
bucketEdge(CLK := btnBucket);
encoderM2(Enable := TRUE, HomingPermit := TRUE, HomingAtTargetM := btnM2 OR bucketEdge.Q, CfgHomingTargetM := 23.7, CfgTopSensorPosM := 23.7, UseDynamicTarget := bucketEdge.Q, DynamicHomingTargetM := encoderM1.Measurement.CablePosM + cfgBucket.OffsetCloseM, HwIn := hw2, Cfg := cfgEncoder, Calib := calibM2); calibM2 := encoderM2.Calib;
bucket(Enable := TRUE, Mode := E_Mode.MAINT_N2, PowerContactorEngaged := TRUE, CablePosM1 := encoderM1.Measurement.CablePosM, CablePosM2 := encoderM2.Measurement.CablePosM, HomedM1 := encoderM1.Homed, HomedM2 := encoderM2.Homed, HomedAndReliableM1 := encoderM1.HomedAndReliable, HomedAndReliableM2 := encoderM2.HomedAndReliable, HomingSuspectM1 := encoderM1.HomingSuspect, HomingSuspectM2 := encoderM2.HomingSuspect, ConfirmClosePosition := btnBucket, Config := cfgBucket, BucketState := bucketState); bucketState := bucket.BucketState;
home.M1Status.HomedAndReliable := encoderM1.HomedAndReliable; home.M2Status.HomedAndReliable := encoderM2.HomedAndReliable; home(BucketOffsetValid := bucketState.BucketReferenced, BtnValidation := bench.Operator.JoyBtnRaw);
ADVANCE_TIME(10000000);
bench(M1_PresetTriggerCmd := encoderM1.HwOut.PresetTriggerCmd, M1_PresetValueOut := encoderM1.HwOut.PresetValueOut, M2_PresetTriggerCmd := encoderM2.HwOut.PresetTriggerCmd, M2_PresetValueOut := encoderM2.HwOut.PresetValueOut, RawPosM1 := raw1, RawPosM2 := raw2); raw1 := bench.RawPosM1; raw2 := bench.RawPosM2;
hw1.RawPosIn := bench.Winch.COD1_PosValue; hw1.SlaveOperational := TRUE; hw2.RawPosIn := bench.Winch.COD2_PosValue; hw2.SlaveOperational := TRUE;
encoderM1(Enable := TRUE, HomingPermit := TRUE, HomingAtTargetM := btnM1, CfgHomingTargetM := 8.7, CfgTopSensorPosM := 8.7, HwIn := hw1, Cfg := cfgEncoder, Calib := calibM1); calibM1 := encoderM1.Calib;
bucketEdge(CLK := btnBucket);
encoderM2(Enable := TRUE, HomingPermit := TRUE, HomingAtTargetM := btnM2 OR bucketEdge.Q, CfgHomingTargetM := 23.7, CfgTopSensorPosM := 23.7, UseDynamicTarget := bucketEdge.Q, DynamicHomingTargetM := encoderM1.Measurement.CablePosM + cfgBucket.OffsetCloseM, HwIn := hw2, Cfg := cfgEncoder, Calib := calibM2); calibM2 := encoderM2.Calib;
bucket(Enable := TRUE, Mode := E_Mode.MAINT_N2, PowerContactorEngaged := TRUE, CablePosM1 := encoderM1.Measurement.CablePosM, CablePosM2 := encoderM2.Measurement.CablePosM, HomedM1 := encoderM1.Homed, HomedM2 := encoderM2.Homed, HomedAndReliableM1 := encoderM1.HomedAndReliable, HomedAndReliableM2 := encoderM2.HomedAndReliable, HomingSuspectM1 := encoderM1.HomingSuspect, HomingSuspectM2 := encoderM2.HomingSuspect, ConfirmClosePosition := btnBucket, Config := cfgBucket, BucketState := bucketState); bucketState := bucket.BucketState;
home.M1Status.HomedAndReliable := encoderM1.HomedAndReliable; home.M2Status.HomedAndReliable := encoderM2.HomedAndReliable; home(BucketOffsetValid := bucketState.BucketReferenced, BtnValidation := bench.Operator.JoyBtnRaw);
ADVANCE_TIME(10000000);
bench(M1_PresetTriggerCmd := encoderM1.HwOut.PresetTriggerCmd, M1_PresetValueOut := encoderM1.HwOut.PresetValueOut, M2_PresetTriggerCmd := encoderM2.HwOut.PresetTriggerCmd, M2_PresetValueOut := encoderM2.HwOut.PresetValueOut, RawPosM1 := raw1, RawPosM2 := raw2); raw1 := bench.RawPosM1; raw2 := bench.RawPosM2;
hw1.RawPosIn := bench.Winch.COD1_PosValue; hw1.SlaveOperational := TRUE; hw2.RawPosIn := bench.Winch.COD2_PosValue; hw2.SlaveOperational := TRUE;
encoderM1(Enable := TRUE, HomingPermit := TRUE, HomingAtTargetM := btnM1, CfgHomingTargetM := 8.7, CfgTopSensorPosM := 8.7, HwIn := hw1, Cfg := cfgEncoder, Calib := calibM1); calibM1 := encoderM1.Calib;
bucketEdge(CLK := btnBucket);
encoderM2(Enable := TRUE, HomingPermit := TRUE, HomingAtTargetM := btnM2 OR bucketEdge.Q, CfgHomingTargetM := 23.7, CfgTopSensorPosM := 23.7, UseDynamicTarget := bucketEdge.Q, DynamicHomingTargetM := encoderM1.Measurement.CablePosM + cfgBucket.OffsetCloseM, HwIn := hw2, Cfg := cfgEncoder, Calib := calibM2); calibM2 := encoderM2.Calib;
bucket(Enable := TRUE, Mode := E_Mode.MAINT_N2, PowerContactorEngaged := TRUE, CablePosM1 := encoderM1.Measurement.CablePosM, CablePosM2 := encoderM2.Measurement.CablePosM, HomedM1 := encoderM1.Homed, HomedM2 := encoderM2.Homed, HomedAndReliableM1 := encoderM1.HomedAndReliable, HomedAndReliableM2 := encoderM2.HomedAndReliable, HomingSuspectM1 := encoderM1.HomingSuspect, HomingSuspectM2 := encoderM2.HomingSuspect, ConfirmClosePosition := btnBucket, Config := cfgBucket, BucketState := bucketState); bucketState := bucket.BucketState;
home.M1Status.HomedAndReliable := encoderM1.HomedAndReliable; home.M2Status.HomedAndReliable := encoderM2.HomedAndReliable; home(BucketOffsetValid := bucketState.BucketReferenced, BtnValidation := bench.Operator.JoyBtnRaw);
ADVANCE_TIME(10000000);
bench(M1_PresetTriggerCmd := encoderM1.HwOut.PresetTriggerCmd, M1_PresetValueOut := encoderM1.HwOut.PresetValueOut, M2_PresetTriggerCmd := encoderM2.HwOut.PresetTriggerCmd, M2_PresetValueOut := encoderM2.HwOut.PresetValueOut, RawPosM1 := raw1, RawPosM2 := raw2); raw1 := bench.RawPosM1; raw2 := bench.RawPosM2;
hw1.RawPosIn := bench.Winch.COD1_PosValue; hw1.SlaveOperational := TRUE; hw2.RawPosIn := bench.Winch.COD2_PosValue; hw2.SlaveOperational := TRUE;
encoderM1(Enable := TRUE, HomingPermit := TRUE, HomingAtTargetM := btnM1, CfgHomingTargetM := 8.7, CfgTopSensorPosM := 8.7, HwIn := hw1, Cfg := cfgEncoder, Calib := calibM1); calibM1 := encoderM1.Calib;
bucketEdge(CLK := btnBucket);
encoderM2(Enable := TRUE, HomingPermit := TRUE, HomingAtTargetM := btnM2 OR bucketEdge.Q, CfgHomingTargetM := 23.7, CfgTopSensorPosM := 23.7, UseDynamicTarget := bucketEdge.Q, DynamicHomingTargetM := encoderM1.Measurement.CablePosM + cfgBucket.OffsetCloseM, HwIn := hw2, Cfg := cfgEncoder, Calib := calibM2); calibM2 := encoderM2.Calib;
bucket(Enable := TRUE, Mode := E_Mode.MAINT_N2, PowerContactorEngaged := TRUE, CablePosM1 := encoderM1.Measurement.CablePosM, CablePosM2 := encoderM2.Measurement.CablePosM, HomedM1 := encoderM1.Homed, HomedM2 := encoderM2.Homed, HomedAndReliableM1 := encoderM1.HomedAndReliable, HomedAndReliableM2 := encoderM2.HomedAndReliable, HomingSuspectM1 := encoderM1.HomingSuspect, HomingSuspectM2 := encoderM2.HomingSuspect, ConfirmClosePosition := btnBucket, Config := cfgBucket, BucketState := bucketState); bucketState := bucket.BucketState;
home.M1Status.HomedAndReliable := encoderM1.HomedAndReliable; home.M2Status.HomedAndReliable := encoderM2.HomedAndReliable; home(BucketOffsetValid := bucketState.BucketReferenced, BtnValidation := bench.Operator.JoyBtnRaw);
ADVANCE_TIME(10000000);
bench(M1_PresetTriggerCmd := encoderM1.HwOut.PresetTriggerCmd, M1_PresetValueOut := encoderM1.HwOut.PresetValueOut, M2_PresetTriggerCmd := encoderM2.HwOut.PresetTriggerCmd, M2_PresetValueOut := encoderM2.HwOut.PresetValueOut, RawPosM1 := raw1, RawPosM2 := raw2); raw1 := bench.RawPosM1; raw2 := bench.RawPosM2;
hw1.RawPosIn := bench.Winch.COD1_PosValue; hw1.SlaveOperational := TRUE; hw2.RawPosIn := bench.Winch.COD2_PosValue; hw2.SlaveOperational := TRUE;
encoderM1(Enable := TRUE, HomingPermit := TRUE, HomingAtTargetM := btnM1, CfgHomingTargetM := 8.7, CfgTopSensorPosM := 8.7, HwIn := hw1, Cfg := cfgEncoder, Calib := calibM1); calibM1 := encoderM1.Calib;
bucketEdge(CLK := btnBucket);
encoderM2(Enable := TRUE, HomingPermit := TRUE, HomingAtTargetM := btnM2 OR bucketEdge.Q, CfgHomingTargetM := 23.7, CfgTopSensorPosM := 23.7, UseDynamicTarget := bucketEdge.Q, DynamicHomingTargetM := encoderM1.Measurement.CablePosM + cfgBucket.OffsetCloseM, HwIn := hw2, Cfg := cfgEncoder, Calib := calibM2); calibM2 := encoderM2.Calib;
bucket(Enable := TRUE, Mode := E_Mode.MAINT_N2, PowerContactorEngaged := TRUE, CablePosM1 := encoderM1.Measurement.CablePosM, CablePosM2 := encoderM2.Measurement.CablePosM, HomedM1 := encoderM1.Homed, HomedM2 := encoderM2.Homed, HomedAndReliableM1 := encoderM1.HomedAndReliable, HomedAndReliableM2 := encoderM2.HomedAndReliable, HomingSuspectM1 := encoderM1.HomingSuspect, HomingSuspectM2 := encoderM2.HomingSuspect, ConfirmClosePosition := btnBucket, Config := cfgBucket, BucketState := bucketState); bucketState := bucket.BucketState;
home.M1Status.HomedAndReliable := encoderM1.HomedAndReliable; home.M2Status.HomedAndReliable := encoderM2.HomedAndReliable; home(BucketOffsetValid := bucketState.BucketReferenced, BtnValidation := bench.Operator.JoyBtnRaw);
ADVANCE_TIME(10000000);
bench(M1_PresetTriggerCmd := encoderM1.HwOut.PresetTriggerCmd, M1_PresetValueOut := encoderM1.HwOut.PresetValueOut, M2_PresetTriggerCmd := encoderM2.HwOut.PresetTriggerCmd, M2_PresetValueOut := encoderM2.HwOut.PresetValueOut, RawPosM1 := raw1, RawPosM2 := raw2); raw1 := bench.RawPosM1; raw2 := bench.RawPosM2;
hw1.RawPosIn := bench.Winch.COD1_PosValue; hw1.SlaveOperational := TRUE; hw2.RawPosIn := bench.Winch.COD2_PosValue; hw2.SlaveOperational := TRUE;
encoderM1(Enable := TRUE, HomingPermit := TRUE, HomingAtTargetM := btnM1, CfgHomingTargetM := 8.7, CfgTopSensorPosM := 8.7, HwIn := hw1, Cfg := cfgEncoder, Calib := calibM1); calibM1 := encoderM1.Calib;
bucketEdge(CLK := btnBucket);
encoderM2(Enable := TRUE, HomingPermit := TRUE, HomingAtTargetM := btnM2 OR bucketEdge.Q, CfgHomingTargetM := 23.7, CfgTopSensorPosM := 23.7, UseDynamicTarget := bucketEdge.Q, DynamicHomingTargetM := encoderM1.Measurement.CablePosM + cfgBucket.OffsetCloseM, HwIn := hw2, Cfg := cfgEncoder, Calib := calibM2); calibM2 := encoderM2.Calib;
bucket(Enable := TRUE, Mode := E_Mode.MAINT_N2, PowerContactorEngaged := TRUE, CablePosM1 := encoderM1.Measurement.CablePosM, CablePosM2 := encoderM2.Measurement.CablePosM, HomedM1 := encoderM1.Homed, HomedM2 := encoderM2.Homed, HomedAndReliableM1 := encoderM1.HomedAndReliable, HomedAndReliableM2 := encoderM2.HomedAndReliable, HomingSuspectM1 := encoderM1.HomingSuspect, HomingSuspectM2 := encoderM2.HomingSuspect, ConfirmClosePosition := btnBucket, Config := cfgBucket, BucketState := bucketState); bucketState := bucket.BucketState;
home.M1Status.HomedAndReliable := encoderM1.HomedAndReliable; home.M2Status.HomedAndReliable := encoderM2.HomedAndReliable; home(BucketOffsetValid := bucketState.BucketReferenced, BtnValidation := bench.Operator.JoyBtnRaw);
ADVANCE_TIME(10000000);
bench(M1_PresetTriggerCmd := encoderM1.HwOut.PresetTriggerCmd, M1_PresetValueOut := encoderM1.HwOut.PresetValueOut, M2_PresetTriggerCmd := encoderM2.HwOut.PresetTriggerCmd, M2_PresetValueOut := encoderM2.HwOut.PresetValueOut, RawPosM1 := raw1, RawPosM2 := raw2); raw1 := bench.RawPosM1; raw2 := bench.RawPosM2;
hw1.RawPosIn := bench.Winch.COD1_PosValue; hw1.SlaveOperational := TRUE; hw2.RawPosIn := bench.Winch.COD2_PosValue; hw2.SlaveOperational := TRUE;
encoderM1(Enable := TRUE, HomingPermit := TRUE, HomingAtTargetM := btnM1, CfgHomingTargetM := 8.7, CfgTopSensorPosM := 8.7, HwIn := hw1, Cfg := cfgEncoder, Calib := calibM1); calibM1 := encoderM1.Calib;
bucketEdge(CLK := btnBucket);
encoderM2(Enable := TRUE, HomingPermit := TRUE, HomingAtTargetM := btnM2 OR bucketEdge.Q, CfgHomingTargetM := 23.7, CfgTopSensorPosM := 23.7, UseDynamicTarget := bucketEdge.Q, DynamicHomingTargetM := encoderM1.Measurement.CablePosM + cfgBucket.OffsetCloseM, HwIn := hw2, Cfg := cfgEncoder, Calib := calibM2); calibM2 := encoderM2.Calib;
bucket(Enable := TRUE, Mode := E_Mode.MAINT_N2, PowerContactorEngaged := TRUE, CablePosM1 := encoderM1.Measurement.CablePosM, CablePosM2 := encoderM2.Measurement.CablePosM, HomedM1 := encoderM1.Homed, HomedM2 := encoderM2.Homed, HomedAndReliableM1 := encoderM1.HomedAndReliable, HomedAndReliableM2 := encoderM2.HomedAndReliable, HomingSuspectM1 := encoderM1.HomingSuspect, HomingSuspectM2 := encoderM2.HomingSuspect, ConfirmClosePosition := btnBucket, Config := cfgBucket, BucketState := bucketState); bucketState := bucket.BucketState;
home.M1Status.HomedAndReliable := encoderM1.HomedAndReliable; home.M2Status.HomedAndReliable := encoderM2.HomedAndReliable; home(BucketOffsetValid := bucketState.BucketReferenced, BtnValidation := bench.Operator.JoyBtnRaw);
ADVANCE_TIME(10000000);
bench(M1_PresetTriggerCmd := encoderM1.HwOut.PresetTriggerCmd, M1_PresetValueOut := encoderM1.HwOut.PresetValueOut, M2_PresetTriggerCmd := encoderM2.HwOut.PresetTriggerCmd, M2_PresetValueOut := encoderM2.HwOut.PresetValueOut, RawPosM1 := raw1, RawPosM2 := raw2); raw1 := bench.RawPosM1; raw2 := bench.RawPosM2;
hw1.RawPosIn := bench.Winch.COD1_PosValue; hw1.SlaveOperational := TRUE; hw2.RawPosIn := bench.Winch.COD2_PosValue; hw2.SlaveOperational := TRUE;
encoderM1(Enable := TRUE, HomingPermit := TRUE, HomingAtTargetM := btnM1, CfgHomingTargetM := 8.7, CfgTopSensorPosM := 8.7, HwIn := hw1, Cfg := cfgEncoder, Calib := calibM1); calibM1 := encoderM1.Calib;
bucketEdge(CLK := btnBucket);
encoderM2(Enable := TRUE, HomingPermit := TRUE, HomingAtTargetM := btnM2 OR bucketEdge.Q, CfgHomingTargetM := 23.7, CfgTopSensorPosM := 23.7, UseDynamicTarget := bucketEdge.Q, DynamicHomingTargetM := encoderM1.Measurement.CablePosM + cfgBucket.OffsetCloseM, HwIn := hw2, Cfg := cfgEncoder, Calib := calibM2); calibM2 := encoderM2.Calib;
bucket(Enable := TRUE, Mode := E_Mode.MAINT_N2, PowerContactorEngaged := TRUE, CablePosM1 := encoderM1.Measurement.CablePosM, CablePosM2 := encoderM2.Measurement.CablePosM, HomedM1 := encoderM1.Homed, HomedM2 := encoderM2.Homed, HomedAndReliableM1 := encoderM1.HomedAndReliable, HomedAndReliableM2 := encoderM2.HomedAndReliable, HomingSuspectM1 := encoderM1.HomingSuspect, HomingSuspectM2 := encoderM2.HomingSuspect, ConfirmClosePosition := btnBucket, Config := cfgBucket, BucketState := bucketState); bucketState := bucket.BucketState;
home.M1Status.HomedAndReliable := encoderM1.HomedAndReliable; home.M2Status.HomedAndReliable := encoderM2.HomedAndReliable; home(BucketOffsetValid := bucketState.BucketReferenced, BtnValidation := bench.Operator.JoyBtnRaw);
ADVANCE_TIME(10000000);
bench(M1_PresetTriggerCmd := encoderM1.HwOut.PresetTriggerCmd, M1_PresetValueOut := encoderM1.HwOut.PresetValueOut, M2_PresetTriggerCmd := encoderM2.HwOut.PresetTriggerCmd, M2_PresetValueOut := encoderM2.HwOut.PresetValueOut, RawPosM1 := raw1, RawPosM2 := raw2); raw1 := bench.RawPosM1; raw2 := bench.RawPosM2;
hw1.RawPosIn := bench.Winch.COD1_PosValue; hw1.SlaveOperational := TRUE; hw2.RawPosIn := bench.Winch.COD2_PosValue; hw2.SlaveOperational := TRUE;
encoderM1(Enable := TRUE, HomingPermit := TRUE, HomingAtTargetM := btnM1, CfgHomingTargetM := 8.7, CfgTopSensorPosM := 8.7, HwIn := hw1, Cfg := cfgEncoder, Calib := calibM1); calibM1 := encoderM1.Calib;
bucketEdge(CLK := btnBucket);
encoderM2(Enable := TRUE, HomingPermit := TRUE, HomingAtTargetM := btnM2 OR bucketEdge.Q, CfgHomingTargetM := 23.7, CfgTopSensorPosM := 23.7, UseDynamicTarget := bucketEdge.Q, DynamicHomingTargetM := encoderM1.Measurement.CablePosM + cfgBucket.OffsetCloseM, HwIn := hw2, Cfg := cfgEncoder, Calib := calibM2); calibM2 := encoderM2.Calib;
bucket(Enable := TRUE, Mode := E_Mode.MAINT_N2, PowerContactorEngaged := TRUE, CablePosM1 := encoderM1.Measurement.CablePosM, CablePosM2 := encoderM2.Measurement.CablePosM, HomedM1 := encoderM1.Homed, HomedM2 := encoderM2.Homed, HomedAndReliableM1 := encoderM1.HomedAndReliable, HomedAndReliableM2 := encoderM2.HomedAndReliable, HomingSuspectM1 := encoderM1.HomingSuspect, HomingSuspectM2 := encoderM2.HomingSuspect, ConfirmClosePosition := btnBucket, Config := cfgBucket, BucketState := bucketState); bucketState := bucket.BucketState;
home.M1Status.HomedAndReliable := encoderM1.HomedAndReliable; home.M2Status.HomedAndReliable := encoderM2.HomedAndReliable; home(BucketOffsetValid := bucketState.BucketReferenced, BtnValidation := bench.Operator.JoyBtnRaw);
ADVANCE_TIME(10000000);
bench(M1_PresetTriggerCmd := encoderM1.HwOut.PresetTriggerCmd, M1_PresetValueOut := encoderM1.HwOut.PresetValueOut, M2_PresetTriggerCmd := encoderM2.HwOut.PresetTriggerCmd, M2_PresetValueOut := encoderM2.HwOut.PresetValueOut, RawPosM1 := raw1, RawPosM2 := raw2); raw1 := bench.RawPosM1; raw2 := bench.RawPosM2;
hw1.RawPosIn := bench.Winch.COD1_PosValue; hw1.SlaveOperational := TRUE; hw2.RawPosIn := bench.Winch.COD2_PosValue; hw2.SlaveOperational := TRUE;
encoderM1(Enable := TRUE, HomingPermit := TRUE, HomingAtTargetM := btnM1, CfgHomingTargetM := 8.7, CfgTopSensorPosM := 8.7, HwIn := hw1, Cfg := cfgEncoder, Calib := calibM1); calibM1 := encoderM1.Calib;
bucketEdge(CLK := btnBucket);
encoderM2(Enable := TRUE, HomingPermit := TRUE, HomingAtTargetM := btnM2 OR bucketEdge.Q, CfgHomingTargetM := 23.7, CfgTopSensorPosM := 23.7, UseDynamicTarget := bucketEdge.Q, DynamicHomingTargetM := encoderM1.Measurement.CablePosM + cfgBucket.OffsetCloseM, HwIn := hw2, Cfg := cfgEncoder, Calib := calibM2); calibM2 := encoderM2.Calib;
bucket(Enable := TRUE, Mode := E_Mode.MAINT_N2, PowerContactorEngaged := TRUE, CablePosM1 := encoderM1.Measurement.CablePosM, CablePosM2 := encoderM2.Measurement.CablePosM, HomedM1 := encoderM1.Homed, HomedM2 := encoderM2.Homed, HomedAndReliableM1 := encoderM1.HomedAndReliable, HomedAndReliableM2 := encoderM2.HomedAndReliable, HomingSuspectM1 := encoderM1.HomingSuspect, HomingSuspectM2 := encoderM2.HomingSuspect, ConfirmClosePosition := btnBucket, Config := cfgBucket, BucketState := bucketState); bucketState := bucket.BucketState;
home.M1Status.HomedAndReliable := encoderM1.HomedAndReliable; home.M2Status.HomedAndReliable := encoderM2.HomedAndReliable; home(BucketOffsetValid := bucketState.BucketReferenced, BtnValidation := bench.Operator.JoyBtnRaw);
ADVANCE_TIME(10000000);
bench(M1_PresetTriggerCmd := encoderM1.HwOut.PresetTriggerCmd, M1_PresetValueOut := encoderM1.HwOut.PresetValueOut, M2_PresetTriggerCmd := encoderM2.HwOut.PresetTriggerCmd, M2_PresetValueOut := encoderM2.HwOut.PresetValueOut, RawPosM1 := raw1, RawPosM2 := raw2); raw1 := bench.RawPosM1; raw2 := bench.RawPosM2;
hw1.RawPosIn := bench.Winch.COD1_PosValue; hw1.SlaveOperational := TRUE; hw2.RawPosIn := bench.Winch.COD2_PosValue; hw2.SlaveOperational := TRUE;
encoderM1(Enable := TRUE, HomingPermit := TRUE, HomingAtTargetM := btnM1, CfgHomingTargetM := 8.7, CfgTopSensorPosM := 8.7, HwIn := hw1, Cfg := cfgEncoder, Calib := calibM1); calibM1 := encoderM1.Calib;
bucketEdge(CLK := btnBucket);
encoderM2(Enable := TRUE, HomingPermit := TRUE, HomingAtTargetM := btnM2 OR bucketEdge.Q, CfgHomingTargetM := 23.7, CfgTopSensorPosM := 23.7, UseDynamicTarget := bucketEdge.Q, DynamicHomingTargetM := encoderM1.Measurement.CablePosM + cfgBucket.OffsetCloseM, HwIn := hw2, Cfg := cfgEncoder, Calib := calibM2); calibM2 := encoderM2.Calib;
bucket(Enable := TRUE, Mode := E_Mode.MAINT_N2, PowerContactorEngaged := TRUE, CablePosM1 := encoderM1.Measurement.CablePosM, CablePosM2 := encoderM2.Measurement.CablePosM, HomedM1 := encoderM1.Homed, HomedM2 := encoderM2.Homed, HomedAndReliableM1 := encoderM1.HomedAndReliable, HomedAndReliableM2 := encoderM2.HomedAndReliable, HomingSuspectM1 := encoderM1.HomingSuspect, HomingSuspectM2 := encoderM2.HomingSuspect, ConfirmClosePosition := btnBucket, Config := cfgBucket, BucketState := bucketState); bucketState := bucket.BucketState;
home.M1Status.HomedAndReliable := encoderM1.HomedAndReliable; home.M2Status.HomedAndReliable := encoderM2.HomedAndReliable; home(BucketOffsetValid := bucketState.BucketReferenced, BtnValidation := bench.Operator.JoyBtnRaw);
ADVANCE_TIME(10000000);
bench(M1_PresetTriggerCmd := encoderM1.HwOut.PresetTriggerCmd, M1_PresetValueOut := encoderM1.HwOut.PresetValueOut, M2_PresetTriggerCmd := encoderM2.HwOut.PresetTriggerCmd, M2_PresetValueOut := encoderM2.HwOut.PresetValueOut, RawPosM1 := raw1, RawPosM2 := raw2); raw1 := bench.RawPosM1; raw2 := bench.RawPosM2;
hw1.RawPosIn := bench.Winch.COD1_PosValue; hw1.SlaveOperational := TRUE; hw2.RawPosIn := bench.Winch.COD2_PosValue; hw2.SlaveOperational := TRUE;
encoderM1(Enable := TRUE, HomingPermit := TRUE, HomingAtTargetM := btnM1, CfgHomingTargetM := 8.7, CfgTopSensorPosM := 8.7, HwIn := hw1, Cfg := cfgEncoder, Calib := calibM1); calibM1 := encoderM1.Calib;
bucketEdge(CLK := btnBucket);
encoderM2(Enable := TRUE, HomingPermit := TRUE, HomingAtTargetM := btnM2 OR bucketEdge.Q, CfgHomingTargetM := 23.7, CfgTopSensorPosM := 23.7, UseDynamicTarget := bucketEdge.Q, DynamicHomingTargetM := encoderM1.Measurement.CablePosM + cfgBucket.OffsetCloseM, HwIn := hw2, Cfg := cfgEncoder, Calib := calibM2); calibM2 := encoderM2.Calib;
bucket(Enable := TRUE, Mode := E_Mode.MAINT_N2, PowerContactorEngaged := TRUE, CablePosM1 := encoderM1.Measurement.CablePosM, CablePosM2 := encoderM2.Measurement.CablePosM, HomedM1 := encoderM1.Homed, HomedM2 := encoderM2.Homed, HomedAndReliableM1 := encoderM1.HomedAndReliable, HomedAndReliableM2 := encoderM2.HomedAndReliable, HomingSuspectM1 := encoderM1.HomingSuspect, HomingSuspectM2 := encoderM2.HomingSuspect, ConfirmClosePosition := btnBucket, Config := cfgBucket, BucketState := bucketState); bucketState := bucket.BucketState;
home.M1Status.HomedAndReliable := encoderM1.HomedAndReliable; home.M2Status.HomedAndReliable := encoderM2.HomedAndReliable; home(BucketOffsetValid := bucketState.BucketReferenced, BtnValidation := bench.Operator.JoyBtnRaw);
ADVANCE_TIME(10000000);
bench(M1_PresetTriggerCmd := encoderM1.HwOut.PresetTriggerCmd, M1_PresetValueOut := encoderM1.HwOut.PresetValueOut, M2_PresetTriggerCmd := encoderM2.HwOut.PresetTriggerCmd, M2_PresetValueOut := encoderM2.HwOut.PresetValueOut, RawPosM1 := raw1, RawPosM2 := raw2); raw1 := bench.RawPosM1; raw2 := bench.RawPosM2;
hw1.RawPosIn := bench.Winch.COD1_PosValue; hw1.SlaveOperational := TRUE; hw2.RawPosIn := bench.Winch.COD2_PosValue; hw2.SlaveOperational := TRUE;
encoderM1(Enable := TRUE, HomingPermit := TRUE, HomingAtTargetM := btnM1, CfgHomingTargetM := 8.7, CfgTopSensorPosM := 8.7, HwIn := hw1, Cfg := cfgEncoder, Calib := calibM1); calibM1 := encoderM1.Calib;
bucketEdge(CLK := btnBucket);
encoderM2(Enable := TRUE, HomingPermit := TRUE, HomingAtTargetM := btnM2 OR bucketEdge.Q, CfgHomingTargetM := 23.7, CfgTopSensorPosM := 23.7, UseDynamicTarget := bucketEdge.Q, DynamicHomingTargetM := encoderM1.Measurement.CablePosM + cfgBucket.OffsetCloseM, HwIn := hw2, Cfg := cfgEncoder, Calib := calibM2); calibM2 := encoderM2.Calib;
bucket(Enable := TRUE, Mode := E_Mode.MAINT_N2, PowerContactorEngaged := TRUE, CablePosM1 := encoderM1.Measurement.CablePosM, CablePosM2 := encoderM2.Measurement.CablePosM, HomedM1 := encoderM1.Homed, HomedM2 := encoderM2.Homed, HomedAndReliableM1 := encoderM1.HomedAndReliable, HomedAndReliableM2 := encoderM2.HomedAndReliable, HomingSuspectM1 := encoderM1.HomingSuspect, HomingSuspectM2 := encoderM2.HomingSuspect, ConfirmClosePosition := btnBucket, Config := cfgBucket, BucketState := bucketState); bucketState := bucket.BucketState;
home.M1Status.HomedAndReliable := encoderM1.HomedAndReliable; home.M2Status.HomedAndReliable := encoderM2.HomedAndReliable; home(BucketOffsetValid := bucketState.BucketReferenced, BtnValidation := bench.Operator.JoyBtnRaw);
ADVANCE_TIME(10000000);
bench(M1_PresetTriggerCmd := encoderM1.HwOut.PresetTriggerCmd, M1_PresetValueOut := encoderM1.HwOut.PresetValueOut, M2_PresetTriggerCmd := encoderM2.HwOut.PresetTriggerCmd, M2_PresetValueOut := encoderM2.HwOut.PresetValueOut, RawPosM1 := raw1, RawPosM2 := raw2); raw1 := bench.RawPosM1; raw2 := bench.RawPosM2;
hw1.RawPosIn := bench.Winch.COD1_PosValue; hw1.SlaveOperational := TRUE; hw2.RawPosIn := bench.Winch.COD2_PosValue; hw2.SlaveOperational := TRUE;
encoderM1(Enable := TRUE, HomingPermit := TRUE, HomingAtTargetM := btnM1, CfgHomingTargetM := 8.7, CfgTopSensorPosM := 8.7, HwIn := hw1, Cfg := cfgEncoder, Calib := calibM1); calibM1 := encoderM1.Calib;
bucketEdge(CLK := btnBucket);
encoderM2(Enable := TRUE, HomingPermit := TRUE, HomingAtTargetM := btnM2 OR bucketEdge.Q, CfgHomingTargetM := 23.7, CfgTopSensorPosM := 23.7, UseDynamicTarget := bucketEdge.Q, DynamicHomingTargetM := encoderM1.Measurement.CablePosM + cfgBucket.OffsetCloseM, HwIn := hw2, Cfg := cfgEncoder, Calib := calibM2); calibM2 := encoderM2.Calib;
bucket(Enable := TRUE, Mode := E_Mode.MAINT_N2, PowerContactorEngaged := TRUE, CablePosM1 := encoderM1.Measurement.CablePosM, CablePosM2 := encoderM2.Measurement.CablePosM, HomedM1 := encoderM1.Homed, HomedM2 := encoderM2.Homed, HomedAndReliableM1 := encoderM1.HomedAndReliable, HomedAndReliableM2 := encoderM2.HomedAndReliable, HomingSuspectM1 := encoderM1.HomingSuspect, HomingSuspectM2 := encoderM2.HomingSuspect, ConfirmClosePosition := btnBucket, Config := cfgBucket, BucketState := bucketState); bucketState := bucket.BucketState;
home.M1Status.HomedAndReliable := encoderM1.HomedAndReliable; home.M2Status.HomedAndReliable := encoderM2.HomedAndReliable; home(BucketOffsetValid := bucketState.BucketReferenced, BtnValidation := bench.Operator.JoyBtnRaw);
ADVANCE_TIME(10000000);
bench(M1_PresetTriggerCmd := encoderM1.HwOut.PresetTriggerCmd, M1_PresetValueOut := encoderM1.HwOut.PresetValueOut, M2_PresetTriggerCmd := encoderM2.HwOut.PresetTriggerCmd, M2_PresetValueOut := encoderM2.HwOut.PresetValueOut, RawPosM1 := raw1, RawPosM2 := raw2); raw1 := bench.RawPosM1; raw2 := bench.RawPosM2;
hw1.RawPosIn := bench.Winch.COD1_PosValue; hw1.SlaveOperational := TRUE; hw2.RawPosIn := bench.Winch.COD2_PosValue; hw2.SlaveOperational := TRUE;
encoderM1(Enable := TRUE, HomingPermit := TRUE, HomingAtTargetM := btnM1, CfgHomingTargetM := 8.7, CfgTopSensorPosM := 8.7, HwIn := hw1, Cfg := cfgEncoder, Calib := calibM1); calibM1 := encoderM1.Calib;
bucketEdge(CLK := btnBucket);
encoderM2(Enable := TRUE, HomingPermit := TRUE, HomingAtTargetM := btnM2 OR bucketEdge.Q, CfgHomingTargetM := 23.7, CfgTopSensorPosM := 23.7, UseDynamicTarget := bucketEdge.Q, DynamicHomingTargetM := encoderM1.Measurement.CablePosM + cfgBucket.OffsetCloseM, HwIn := hw2, Cfg := cfgEncoder, Calib := calibM2); calibM2 := encoderM2.Calib;
bucket(Enable := TRUE, Mode := E_Mode.MAINT_N2, PowerContactorEngaged := TRUE, CablePosM1 := encoderM1.Measurement.CablePosM, CablePosM2 := encoderM2.Measurement.CablePosM, HomedM1 := encoderM1.Homed, HomedM2 := encoderM2.Homed, HomedAndReliableM1 := encoderM1.HomedAndReliable, HomedAndReliableM2 := encoderM2.HomedAndReliable, HomingSuspectM1 := encoderM1.HomingSuspect, HomingSuspectM2 := encoderM2.HomingSuspect, ConfirmClosePosition := btnBucket, Config := cfgBucket, BucketState := bucketState); bucketState := bucket.BucketState;
home.M1Status.HomedAndReliable := encoderM1.HomedAndReliable; home.M2Status.HomedAndReliable := encoderM2.HomedAndReliable; home(BucketOffsetValid := bucketState.BucketReferenced, BtnValidation := bench.Operator.JoyBtnRaw);
ADVANCE_TIME(10000000);
bench(M1_PresetTriggerCmd := encoderM1.HwOut.PresetTriggerCmd, M1_PresetValueOut := encoderM1.HwOut.PresetValueOut, M2_PresetTriggerCmd := encoderM2.HwOut.PresetTriggerCmd, M2_PresetValueOut := encoderM2.HwOut.PresetValueOut, RawPosM1 := raw1, RawPosM2 := raw2); raw1 := bench.RawPosM1; raw2 := bench.RawPosM2;
hw1.RawPosIn := bench.Winch.COD1_PosValue; hw1.SlaveOperational := TRUE; hw2.RawPosIn := bench.Winch.COD2_PosValue; hw2.SlaveOperational := TRUE;
encoderM1(Enable := TRUE, HomingPermit := TRUE, HomingAtTargetM := btnM1, CfgHomingTargetM := 8.7, CfgTopSensorPosM := 8.7, HwIn := hw1, Cfg := cfgEncoder, Calib := calibM1); calibM1 := encoderM1.Calib;
bucketEdge(CLK := btnBucket);
encoderM2(Enable := TRUE, HomingPermit := TRUE, HomingAtTargetM := btnM2 OR bucketEdge.Q, CfgHomingTargetM := 23.7, CfgTopSensorPosM := 23.7, UseDynamicTarget := bucketEdge.Q, DynamicHomingTargetM := encoderM1.Measurement.CablePosM + cfgBucket.OffsetCloseM, HwIn := hw2, Cfg := cfgEncoder, Calib := calibM2); calibM2 := encoderM2.Calib;
bucket(Enable := TRUE, Mode := E_Mode.MAINT_N2, PowerContactorEngaged := TRUE, CablePosM1 := encoderM1.Measurement.CablePosM, CablePosM2 := encoderM2.Measurement.CablePosM, HomedM1 := encoderM1.Homed, HomedM2 := encoderM2.Homed, HomedAndReliableM1 := encoderM1.HomedAndReliable, HomedAndReliableM2 := encoderM2.HomedAndReliable, HomingSuspectM1 := encoderM1.HomingSuspect, HomingSuspectM2 := encoderM2.HomingSuspect, ConfirmClosePosition := btnBucket, Config := cfgBucket, BucketState := bucketState); bucketState := bucket.BucketState;
home.M1Status.HomedAndReliable := encoderM1.HomedAndReliable; home.M2Status.HomedAndReliable := encoderM2.HomedAndReliable; home(BucketOffsetValid := bucketState.BucketReferenced, BtnValidation := bench.Operator.JoyBtnRaw);
ADVANCE_TIME(10000000);
bench(M1_PresetTriggerCmd := encoderM1.HwOut.PresetTriggerCmd, M1_PresetValueOut := encoderM1.HwOut.PresetValueOut, M2_PresetTriggerCmd := encoderM2.HwOut.PresetTriggerCmd, M2_PresetValueOut := encoderM2.HwOut.PresetValueOut, RawPosM1 := raw1, RawPosM2 := raw2); raw1 := bench.RawPosM1; raw2 := bench.RawPosM2;
hw1.RawPosIn := bench.Winch.COD1_PosValue; hw1.SlaveOperational := TRUE; hw2.RawPosIn := bench.Winch.COD2_PosValue; hw2.SlaveOperational := TRUE;
encoderM1(Enable := TRUE, HomingPermit := TRUE, HomingAtTargetM := btnM1, CfgHomingTargetM := 8.7, CfgTopSensorPosM := 8.7, HwIn := hw1, Cfg := cfgEncoder, Calib := calibM1); calibM1 := encoderM1.Calib;
bucketEdge(CLK := btnBucket);
encoderM2(Enable := TRUE, HomingPermit := TRUE, HomingAtTargetM := btnM2 OR bucketEdge.Q, CfgHomingTargetM := 23.7, CfgTopSensorPosM := 23.7, UseDynamicTarget := bucketEdge.Q, DynamicHomingTargetM := encoderM1.Measurement.CablePosM + cfgBucket.OffsetCloseM, HwIn := hw2, Cfg := cfgEncoder, Calib := calibM2); calibM2 := encoderM2.Calib;
bucket(Enable := TRUE, Mode := E_Mode.MAINT_N2, PowerContactorEngaged := TRUE, CablePosM1 := encoderM1.Measurement.CablePosM, CablePosM2 := encoderM2.Measurement.CablePosM, HomedM1 := encoderM1.Homed, HomedM2 := encoderM2.Homed, HomedAndReliableM1 := encoderM1.HomedAndReliable, HomedAndReliableM2 := encoderM2.HomedAndReliable, HomingSuspectM1 := encoderM1.HomingSuspect, HomingSuspectM2 := encoderM2.HomingSuspect, ConfirmClosePosition := btnBucket, Config := cfgBucket, BucketState := bucketState); bucketState := bucket.BucketState;
home.M1Status.HomedAndReliable := encoderM1.HomedAndReliable; home.M2Status.HomedAndReliable := encoderM2.HomedAndReliable; home(BucketOffsetValid := bucketState.BucketReferenced, BtnValidation := bench.Operator.JoyBtnRaw);
ADVANCE_TIME(10000000);
bench(M1_PresetTriggerCmd := encoderM1.HwOut.PresetTriggerCmd, M1_PresetValueOut := encoderM1.HwOut.PresetValueOut, M2_PresetTriggerCmd := encoderM2.HwOut.PresetTriggerCmd, M2_PresetValueOut := encoderM2.HwOut.PresetValueOut, RawPosM1 := raw1, RawPosM2 := raw2); raw1 := bench.RawPosM1; raw2 := bench.RawPosM2;
hw1.RawPosIn := bench.Winch.COD1_PosValue; hw1.SlaveOperational := TRUE; hw2.RawPosIn := bench.Winch.COD2_PosValue; hw2.SlaveOperational := TRUE;
encoderM1(Enable := TRUE, HomingPermit := TRUE, HomingAtTargetM := btnM1, CfgHomingTargetM := 8.7, CfgTopSensorPosM := 8.7, HwIn := hw1, Cfg := cfgEncoder, Calib := calibM1); calibM1 := encoderM1.Calib;
bucketEdge(CLK := btnBucket);
encoderM2(Enable := TRUE, HomingPermit := TRUE, HomingAtTargetM := btnM2 OR bucketEdge.Q, CfgHomingTargetM := 23.7, CfgTopSensorPosM := 23.7, UseDynamicTarget := bucketEdge.Q, DynamicHomingTargetM := encoderM1.Measurement.CablePosM + cfgBucket.OffsetCloseM, HwIn := hw2, Cfg := cfgEncoder, Calib := calibM2); calibM2 := encoderM2.Calib;
bucket(Enable := TRUE, Mode := E_Mode.MAINT_N2, PowerContactorEngaged := TRUE, CablePosM1 := encoderM1.Measurement.CablePosM, CablePosM2 := encoderM2.Measurement.CablePosM, HomedM1 := encoderM1.Homed, HomedM2 := encoderM2.Homed, HomedAndReliableM1 := encoderM1.HomedAndReliable, HomedAndReliableM2 := encoderM2.HomedAndReliable, HomingSuspectM1 := encoderM1.HomingSuspect, HomingSuspectM2 := encoderM2.HomingSuspect, ConfirmClosePosition := btnBucket, Config := cfgBucket, BucketState := bucketState); bucketState := bucket.BucketState;
home.M1Status.HomedAndReliable := encoderM1.HomedAndReliable; home.M2Status.HomedAndReliable := encoderM2.HomedAndReliable; home(BucketOffsetValid := bucketState.BucketReferenced, BtnValidation := bench.Operator.JoyBtnRaw);
ADVANCE_TIME(10000000);
bench(M1_PresetTriggerCmd := encoderM1.HwOut.PresetTriggerCmd, M1_PresetValueOut := encoderM1.HwOut.PresetValueOut, M2_PresetTriggerCmd := encoderM2.HwOut.PresetTriggerCmd, M2_PresetValueOut := encoderM2.HwOut.PresetValueOut, RawPosM1 := raw1, RawPosM2 := raw2); raw1 := bench.RawPosM1; raw2 := bench.RawPosM2;
hw1.RawPosIn := bench.Winch.COD1_PosValue; hw1.SlaveOperational := TRUE; hw2.RawPosIn := bench.Winch.COD2_PosValue; hw2.SlaveOperational := TRUE;
encoderM1(Enable := TRUE, HomingPermit := TRUE, HomingAtTargetM := btnM1, CfgHomingTargetM := 8.7, CfgTopSensorPosM := 8.7, HwIn := hw1, Cfg := cfgEncoder, Calib := calibM1); calibM1 := encoderM1.Calib;
bucketEdge(CLK := btnBucket);
encoderM2(Enable := TRUE, HomingPermit := TRUE, HomingAtTargetM := btnM2 OR bucketEdge.Q, CfgHomingTargetM := 23.7, CfgTopSensorPosM := 23.7, UseDynamicTarget := bucketEdge.Q, DynamicHomingTargetM := encoderM1.Measurement.CablePosM + cfgBucket.OffsetCloseM, HwIn := hw2, Cfg := cfgEncoder, Calib := calibM2); calibM2 := encoderM2.Calib;
bucket(Enable := TRUE, Mode := E_Mode.MAINT_N2, PowerContactorEngaged := TRUE, CablePosM1 := encoderM1.Measurement.CablePosM, CablePosM2 := encoderM2.Measurement.CablePosM, HomedM1 := encoderM1.Homed, HomedM2 := encoderM2.Homed, HomedAndReliableM1 := encoderM1.HomedAndReliable, HomedAndReliableM2 := encoderM2.HomedAndReliable, HomingSuspectM1 := encoderM1.HomingSuspect, HomingSuspectM2 := encoderM2.HomingSuspect, ConfirmClosePosition := btnBucket, Config := cfgBucket, BucketState := bucketState); bucketState := bucket.BucketState;
home.M1Status.HomedAndReliable := encoderM1.HomedAndReliable; home.M2Status.HomedAndReliable := encoderM2.HomedAndReliable; home(BucketOffsetValid := bucketState.BucketReferenced, BtnValidation := bench.Operator.JoyBtnRaw);
ADVANCE_TIME(10000000);
bench(M1_PresetTriggerCmd := encoderM1.HwOut.PresetTriggerCmd, M1_PresetValueOut := encoderM1.HwOut.PresetValueOut, M2_PresetTriggerCmd := encoderM2.HwOut.PresetTriggerCmd, M2_PresetValueOut := encoderM2.HwOut.PresetValueOut, RawPosM1 := raw1, RawPosM2 := raw2); raw1 := bench.RawPosM1; raw2 := bench.RawPosM2;
hw1.RawPosIn := bench.Winch.COD1_PosValue; hw1.SlaveOperational := TRUE; hw2.RawPosIn := bench.Winch.COD2_PosValue; hw2.SlaveOperational := TRUE;
encoderM1(Enable := TRUE, HomingPermit := TRUE, HomingAtTargetM := btnM1, CfgHomingTargetM := 8.7, CfgTopSensorPosM := 8.7, HwIn := hw1, Cfg := cfgEncoder, Calib := calibM1); calibM1 := encoderM1.Calib;
bucketEdge(CLK := btnBucket);
encoderM2(Enable := TRUE, HomingPermit := TRUE, HomingAtTargetM := btnM2 OR bucketEdge.Q, CfgHomingTargetM := 23.7, CfgTopSensorPosM := 23.7, UseDynamicTarget := bucketEdge.Q, DynamicHomingTargetM := encoderM1.Measurement.CablePosM + cfgBucket.OffsetCloseM, HwIn := hw2, Cfg := cfgEncoder, Calib := calibM2); calibM2 := encoderM2.Calib;
bucket(Enable := TRUE, Mode := E_Mode.MAINT_N2, PowerContactorEngaged := TRUE, CablePosM1 := encoderM1.Measurement.CablePosM, CablePosM2 := encoderM2.Measurement.CablePosM, HomedM1 := encoderM1.Homed, HomedM2 := encoderM2.Homed, HomedAndReliableM1 := encoderM1.HomedAndReliable, HomedAndReliableM2 := encoderM2.HomedAndReliable, HomingSuspectM1 := encoderM1.HomingSuspect, HomingSuspectM2 := encoderM2.HomingSuspect, ConfirmClosePosition := btnBucket, Config := cfgBucket, BucketState := bucketState); bucketState := bucket.BucketState;
home.M1Status.HomedAndReliable := encoderM1.HomedAndReliable; home.M2Status.HomedAndReliable := encoderM2.HomedAndReliable; home(BucketOffsetValid := bucketState.BucketReferenced, BtnValidation := bench.Operator.JoyBtnRaw);
ADVANCE_TIME(10000000);
bench(M1_PresetTriggerCmd := encoderM1.HwOut.PresetTriggerCmd, M1_PresetValueOut := encoderM1.HwOut.PresetValueOut, M2_PresetTriggerCmd := encoderM2.HwOut.PresetTriggerCmd, M2_PresetValueOut := encoderM2.HwOut.PresetValueOut, RawPosM1 := raw1, RawPosM2 := raw2); raw1 := bench.RawPosM1; raw2 := bench.RawPosM2;
hw1.RawPosIn := bench.Winch.COD1_PosValue; hw1.SlaveOperational := TRUE; hw2.RawPosIn := bench.Winch.COD2_PosValue; hw2.SlaveOperational := TRUE;
encoderM1(Enable := TRUE, HomingPermit := TRUE, HomingAtTargetM := btnM1, CfgHomingTargetM := 8.7, CfgTopSensorPosM := 8.7, HwIn := hw1, Cfg := cfgEncoder, Calib := calibM1); calibM1 := encoderM1.Calib;
bucketEdge(CLK := btnBucket);
encoderM2(Enable := TRUE, HomingPermit := TRUE, HomingAtTargetM := btnM2 OR bucketEdge.Q, CfgHomingTargetM := 23.7, CfgTopSensorPosM := 23.7, UseDynamicTarget := bucketEdge.Q, DynamicHomingTargetM := encoderM1.Measurement.CablePosM + cfgBucket.OffsetCloseM, HwIn := hw2, Cfg := cfgEncoder, Calib := calibM2); calibM2 := encoderM2.Calib;
bucket(Enable := TRUE, Mode := E_Mode.MAINT_N2, PowerContactorEngaged := TRUE, CablePosM1 := encoderM1.Measurement.CablePosM, CablePosM2 := encoderM2.Measurement.CablePosM, HomedM1 := encoderM1.Homed, HomedM2 := encoderM2.Homed, HomedAndReliableM1 := encoderM1.HomedAndReliable, HomedAndReliableM2 := encoderM2.HomedAndReliable, HomingSuspectM1 := encoderM1.HomingSuspect, HomingSuspectM2 := encoderM2.HomingSuspect, ConfirmClosePosition := btnBucket, Config := cfgBucket, BucketState := bucketState); bucketState := bucket.BucketState;
home.M1Status.HomedAndReliable := encoderM1.HomedAndReliable; home.M2Status.HomedAndReliable := encoderM2.HomedAndReliable; home(BucketOffsetValid := bucketState.BucketReferenced, BtnValidation := bench.Operator.JoyBtnRaw);
ADVANCE_TIME(10000000);
bench(M1_PresetTriggerCmd := encoderM1.HwOut.PresetTriggerCmd, M1_PresetValueOut := encoderM1.HwOut.PresetValueOut, M2_PresetTriggerCmd := encoderM2.HwOut.PresetTriggerCmd, M2_PresetValueOut := encoderM2.HwOut.PresetValueOut, RawPosM1 := raw1, RawPosM2 := raw2); raw1 := bench.RawPosM1; raw2 := bench.RawPosM2;
hw1.RawPosIn := bench.Winch.COD1_PosValue; hw1.SlaveOperational := TRUE; hw2.RawPosIn := bench.Winch.COD2_PosValue; hw2.SlaveOperational := TRUE;
encoderM1(Enable := TRUE, HomingPermit := TRUE, HomingAtTargetM := btnM1, CfgHomingTargetM := 8.7, CfgTopSensorPosM := 8.7, HwIn := hw1, Cfg := cfgEncoder, Calib := calibM1); calibM1 := encoderM1.Calib;
bucketEdge(CLK := btnBucket);
encoderM2(Enable := TRUE, HomingPermit := TRUE, HomingAtTargetM := btnM2 OR bucketEdge.Q, CfgHomingTargetM := 23.7, CfgTopSensorPosM := 23.7, UseDynamicTarget := bucketEdge.Q, DynamicHomingTargetM := encoderM1.Measurement.CablePosM + cfgBucket.OffsetCloseM, HwIn := hw2, Cfg := cfgEncoder, Calib := calibM2); calibM2 := encoderM2.Calib;
bucket(Enable := TRUE, Mode := E_Mode.MAINT_N2, PowerContactorEngaged := TRUE, CablePosM1 := encoderM1.Measurement.CablePosM, CablePosM2 := encoderM2.Measurement.CablePosM, HomedM1 := encoderM1.Homed, HomedM2 := encoderM2.Homed, HomedAndReliableM1 := encoderM1.HomedAndReliable, HomedAndReliableM2 := encoderM2.HomedAndReliable, HomingSuspectM1 := encoderM1.HomingSuspect, HomingSuspectM2 := encoderM2.HomingSuspect, ConfirmClosePosition := btnBucket, Config := cfgBucket, BucketState := bucketState); bucketState := bucket.BucketState;
home.M1Status.HomedAndReliable := encoderM1.HomedAndReliable; home.M2Status.HomedAndReliable := encoderM2.HomedAndReliable; home(BucketOffsetValid := bucketState.BucketReferenced, BtnValidation := bench.Operator.JoyBtnRaw);
ADVANCE_TIME(10000000);
bench(M1_PresetTriggerCmd := encoderM1.HwOut.PresetTriggerCmd, M1_PresetValueOut := encoderM1.HwOut.PresetValueOut, M2_PresetTriggerCmd := encoderM2.HwOut.PresetTriggerCmd, M2_PresetValueOut := encoderM2.HwOut.PresetValueOut, RawPosM1 := raw1, RawPosM2 := raw2); raw1 := bench.RawPosM1; raw2 := bench.RawPosM2;
hw1.RawPosIn := bench.Winch.COD1_PosValue; hw1.SlaveOperational := TRUE; hw2.RawPosIn := bench.Winch.COD2_PosValue; hw2.SlaveOperational := TRUE;
encoderM1(Enable := TRUE, HomingPermit := TRUE, HomingAtTargetM := btnM1, CfgHomingTargetM := 8.7, CfgTopSensorPosM := 8.7, HwIn := hw1, Cfg := cfgEncoder, Calib := calibM1); calibM1 := encoderM1.Calib;
bucketEdge(CLK := btnBucket);
encoderM2(Enable := TRUE, HomingPermit := TRUE, HomingAtTargetM := btnM2 OR bucketEdge.Q, CfgHomingTargetM := 23.7, CfgTopSensorPosM := 23.7, UseDynamicTarget := bucketEdge.Q, DynamicHomingTargetM := encoderM1.Measurement.CablePosM + cfgBucket.OffsetCloseM, HwIn := hw2, Cfg := cfgEncoder, Calib := calibM2); calibM2 := encoderM2.Calib;
bucket(Enable := TRUE, Mode := E_Mode.MAINT_N2, PowerContactorEngaged := TRUE, CablePosM1 := encoderM1.Measurement.CablePosM, CablePosM2 := encoderM2.Measurement.CablePosM, HomedM1 := encoderM1.Homed, HomedM2 := encoderM2.Homed, HomedAndReliableM1 := encoderM1.HomedAndReliable, HomedAndReliableM2 := encoderM2.HomedAndReliable, HomingSuspectM1 := encoderM1.HomingSuspect, HomingSuspectM2 := encoderM2.HomingSuspect, ConfirmClosePosition := btnBucket, Config := cfgBucket, BucketState := bucketState); bucketState := bucket.BucketState;
home.M1Status.HomedAndReliable := encoderM1.HomedAndReliable; home.M2Status.HomedAndReliable := encoderM2.HomedAndReliable; home(BucketOffsetValid := bucketState.BucketReferenced, BtnValidation := bench.Operator.JoyBtnRaw);
ADVANCE_TIME(10000000);
bench(M1_PresetTriggerCmd := encoderM1.HwOut.PresetTriggerCmd, M1_PresetValueOut := encoderM1.HwOut.PresetValueOut, M2_PresetTriggerCmd := encoderM2.HwOut.PresetTriggerCmd, M2_PresetValueOut := encoderM2.HwOut.PresetValueOut, RawPosM1 := raw1, RawPosM2 := raw2); raw1 := bench.RawPosM1; raw2 := bench.RawPosM2;
hw1.RawPosIn := bench.Winch.COD1_PosValue; hw1.SlaveOperational := TRUE; hw2.RawPosIn := bench.Winch.COD2_PosValue; hw2.SlaveOperational := TRUE;
encoderM1(Enable := TRUE, HomingPermit := TRUE, HomingAtTargetM := btnM1, CfgHomingTargetM := 8.7, CfgTopSensorPosM := 8.7, HwIn := hw1, Cfg := cfgEncoder, Calib := calibM1); calibM1 := encoderM1.Calib;
bucketEdge(CLK := btnBucket);
encoderM2(Enable := TRUE, HomingPermit := TRUE, HomingAtTargetM := btnM2 OR bucketEdge.Q, CfgHomingTargetM := 23.7, CfgTopSensorPosM := 23.7, UseDynamicTarget := bucketEdge.Q, DynamicHomingTargetM := encoderM1.Measurement.CablePosM + cfgBucket.OffsetCloseM, HwIn := hw2, Cfg := cfgEncoder, Calib := calibM2); calibM2 := encoderM2.Calib;
bucket(Enable := TRUE, Mode := E_Mode.MAINT_N2, PowerContactorEngaged := TRUE, CablePosM1 := encoderM1.Measurement.CablePosM, CablePosM2 := encoderM2.Measurement.CablePosM, HomedM1 := encoderM1.Homed, HomedM2 := encoderM2.Homed, HomedAndReliableM1 := encoderM1.HomedAndReliable, HomedAndReliableM2 := encoderM2.HomedAndReliable, HomingSuspectM1 := encoderM1.HomingSuspect, HomingSuspectM2 := encoderM2.HomingSuspect, ConfirmClosePosition := btnBucket, Config := cfgBucket, BucketState := bucketState); bucketState := bucket.BucketState;
home.M1Status.HomedAndReliable := encoderM1.HomedAndReliable; home.M2Status.HomedAndReliable := encoderM2.HomedAndReliable; home(BucketOffsetValid := bucketState.BucketReferenced, BtnValidation := bench.Operator.JoyBtnRaw);
ADVANCE_TIME(10000000);
bench(M1_PresetTriggerCmd := encoderM1.HwOut.PresetTriggerCmd, M1_PresetValueOut := encoderM1.HwOut.PresetValueOut, M2_PresetTriggerCmd := encoderM2.HwOut.PresetTriggerCmd, M2_PresetValueOut := encoderM2.HwOut.PresetValueOut, RawPosM1 := raw1, RawPosM2 := raw2); raw1 := bench.RawPosM1; raw2 := bench.RawPosM2;
hw1.RawPosIn := bench.Winch.COD1_PosValue; hw1.SlaveOperational := TRUE; hw2.RawPosIn := bench.Winch.COD2_PosValue; hw2.SlaveOperational := TRUE;
encoderM1(Enable := TRUE, HomingPermit := TRUE, HomingAtTargetM := btnM1, CfgHomingTargetM := 8.7, CfgTopSensorPosM := 8.7, HwIn := hw1, Cfg := cfgEncoder, Calib := calibM1); calibM1 := encoderM1.Calib;
bucketEdge(CLK := btnBucket);
encoderM2(Enable := TRUE, HomingPermit := TRUE, HomingAtTargetM := btnM2 OR bucketEdge.Q, CfgHomingTargetM := 23.7, CfgTopSensorPosM := 23.7, UseDynamicTarget := bucketEdge.Q, DynamicHomingTargetM := encoderM1.Measurement.CablePosM + cfgBucket.OffsetCloseM, HwIn := hw2, Cfg := cfgEncoder, Calib := calibM2); calibM2 := encoderM2.Calib;
bucket(Enable := TRUE, Mode := E_Mode.MAINT_N2, PowerContactorEngaged := TRUE, CablePosM1 := encoderM1.Measurement.CablePosM, CablePosM2 := encoderM2.Measurement.CablePosM, HomedM1 := encoderM1.Homed, HomedM2 := encoderM2.Homed, HomedAndReliableM1 := encoderM1.HomedAndReliable, HomedAndReliableM2 := encoderM2.HomedAndReliable, HomingSuspectM1 := encoderM1.HomingSuspect, HomingSuspectM2 := encoderM2.HomingSuspect, ConfirmClosePosition := btnBucket, Config := cfgBucket, BucketState := bucketState); bucketState := bucket.BucketState;
home.M1Status.HomedAndReliable := encoderM1.HomedAndReliable; home.M2Status.HomedAndReliable := encoderM2.HomedAndReliable; home(BucketOffsetValid := bucketState.BucketReferenced, BtnValidation := bench.Operator.JoyBtnRaw);
ADVANCE_TIME(10000000);
bench(M1_PresetTriggerCmd := encoderM1.HwOut.PresetTriggerCmd, M1_PresetValueOut := encoderM1.HwOut.PresetValueOut, M2_PresetTriggerCmd := encoderM2.HwOut.PresetTriggerCmd, M2_PresetValueOut := encoderM2.HwOut.PresetValueOut, RawPosM1 := raw1, RawPosM2 := raw2); raw1 := bench.RawPosM1; raw2 := bench.RawPosM2;
hw1.RawPosIn := bench.Winch.COD1_PosValue; hw1.SlaveOperational := TRUE; hw2.RawPosIn := bench.Winch.COD2_PosValue; hw2.SlaveOperational := TRUE;
encoderM1(Enable := TRUE, HomingPermit := TRUE, HomingAtTargetM := btnM1, CfgHomingTargetM := 8.7, CfgTopSensorPosM := 8.7, HwIn := hw1, Cfg := cfgEncoder, Calib := calibM1); calibM1 := encoderM1.Calib;
bucketEdge(CLK := btnBucket);
encoderM2(Enable := TRUE, HomingPermit := TRUE, HomingAtTargetM := btnM2 OR bucketEdge.Q, CfgHomingTargetM := 23.7, CfgTopSensorPosM := 23.7, UseDynamicTarget := bucketEdge.Q, DynamicHomingTargetM := encoderM1.Measurement.CablePosM + cfgBucket.OffsetCloseM, HwIn := hw2, Cfg := cfgEncoder, Calib := calibM2); calibM2 := encoderM2.Calib;
bucket(Enable := TRUE, Mode := E_Mode.MAINT_N2, PowerContactorEngaged := TRUE, CablePosM1 := encoderM1.Measurement.CablePosM, CablePosM2 := encoderM2.Measurement.CablePosM, HomedM1 := encoderM1.Homed, HomedM2 := encoderM2.Homed, HomedAndReliableM1 := encoderM1.HomedAndReliable, HomedAndReliableM2 := encoderM2.HomedAndReliable, HomingSuspectM1 := encoderM1.HomingSuspect, HomingSuspectM2 := encoderM2.HomingSuspect, ConfirmClosePosition := btnBucket, Config := cfgBucket, BucketState := bucketState); bucketState := bucket.BucketState;
home.M1Status.HomedAndReliable := encoderM1.HomedAndReliable; home.M2Status.HomedAndReliable := encoderM2.HomedAndReliable; home(BucketOffsetValid := bucketState.BucketReferenced, BtnValidation := bench.Operator.JoyBtnRaw);
ADVANCE_TIME(10000000);
bench(M1_PresetTriggerCmd := encoderM1.HwOut.PresetTriggerCmd, M1_PresetValueOut := encoderM1.HwOut.PresetValueOut, M2_PresetTriggerCmd := encoderM2.HwOut.PresetTriggerCmd, M2_PresetValueOut := encoderM2.HwOut.PresetValueOut, RawPosM1 := raw1, RawPosM2 := raw2); raw1 := bench.RawPosM1; raw2 := bench.RawPosM2;
hw1.RawPosIn := bench.Winch.COD1_PosValue; hw1.SlaveOperational := TRUE; hw2.RawPosIn := bench.Winch.COD2_PosValue; hw2.SlaveOperational := TRUE;
encoderM1(Enable := TRUE, HomingPermit := TRUE, HomingAtTargetM := btnM1, CfgHomingTargetM := 8.7, CfgTopSensorPosM := 8.7, HwIn := hw1, Cfg := cfgEncoder, Calib := calibM1); calibM1 := encoderM1.Calib;
bucketEdge(CLK := btnBucket);
encoderM2(Enable := TRUE, HomingPermit := TRUE, HomingAtTargetM := btnM2 OR bucketEdge.Q, CfgHomingTargetM := 23.7, CfgTopSensorPosM := 23.7, UseDynamicTarget := bucketEdge.Q, DynamicHomingTargetM := encoderM1.Measurement.CablePosM + cfgBucket.OffsetCloseM, HwIn := hw2, Cfg := cfgEncoder, Calib := calibM2); calibM2 := encoderM2.Calib;
bucket(Enable := TRUE, Mode := E_Mode.MAINT_N2, PowerContactorEngaged := TRUE, CablePosM1 := encoderM1.Measurement.CablePosM, CablePosM2 := encoderM2.Measurement.CablePosM, HomedM1 := encoderM1.Homed, HomedM2 := encoderM2.Homed, HomedAndReliableM1 := encoderM1.HomedAndReliable, HomedAndReliableM2 := encoderM2.HomedAndReliable, HomingSuspectM1 := encoderM1.HomingSuspect, HomingSuspectM2 := encoderM2.HomingSuspect, ConfirmClosePosition := btnBucket, Config := cfgBucket, BucketState := bucketState); bucketState := bucket.BucketState;
home.M1Status.HomedAndReliable := encoderM1.HomedAndReliable; home.M2Status.HomedAndReliable := encoderM2.HomedAndReliable; home(BucketOffsetValid := bucketState.BucketReferenced, BtnValidation := bench.Operator.JoyBtnRaw);
ADVANCE_TIME(10000000);
bench(M1_PresetTriggerCmd := encoderM1.HwOut.PresetTriggerCmd, M1_PresetValueOut := encoderM1.HwOut.PresetValueOut, M2_PresetTriggerCmd := encoderM2.HwOut.PresetTriggerCmd, M2_PresetValueOut := encoderM2.HwOut.PresetValueOut, RawPosM1 := raw1, RawPosM2 := raw2); raw1 := bench.RawPosM1; raw2 := bench.RawPosM2;
hw1.RawPosIn := bench.Winch.COD1_PosValue; hw1.SlaveOperational := TRUE; hw2.RawPosIn := bench.Winch.COD2_PosValue; hw2.SlaveOperational := TRUE;
encoderM1(Enable := TRUE, HomingPermit := TRUE, HomingAtTargetM := btnM1, CfgHomingTargetM := 8.7, CfgTopSensorPosM := 8.7, HwIn := hw1, Cfg := cfgEncoder, Calib := calibM1); calibM1 := encoderM1.Calib;
bucketEdge(CLK := btnBucket);
encoderM2(Enable := TRUE, HomingPermit := TRUE, HomingAtTargetM := btnM2 OR bucketEdge.Q, CfgHomingTargetM := 23.7, CfgTopSensorPosM := 23.7, UseDynamicTarget := bucketEdge.Q, DynamicHomingTargetM := encoderM1.Measurement.CablePosM + cfgBucket.OffsetCloseM, HwIn := hw2, Cfg := cfgEncoder, Calib := calibM2); calibM2 := encoderM2.Calib;
bucket(Enable := TRUE, Mode := E_Mode.MAINT_N2, PowerContactorEngaged := TRUE, CablePosM1 := encoderM1.Measurement.CablePosM, CablePosM2 := encoderM2.Measurement.CablePosM, HomedM1 := encoderM1.Homed, HomedM2 := encoderM2.Homed, HomedAndReliableM1 := encoderM1.HomedAndReliable, HomedAndReliableM2 := encoderM2.HomedAndReliable, HomingSuspectM1 := encoderM1.HomingSuspect, HomingSuspectM2 := encoderM2.HomingSuspect, ConfirmClosePosition := btnBucket, Config := cfgBucket, BucketState := bucketState); bucketState := bucket.BucketState;
home.M1Status.HomedAndReliable := encoderM1.HomedAndReliable; home.M2Status.HomedAndReliable := encoderM2.HomedAndReliable; home(BucketOffsetValid := bucketState.BucketReferenced, BtnValidation := bench.Operator.JoyBtnRaw);
ADVANCE_TIME(10000000);
bench(M1_PresetTriggerCmd := encoderM1.HwOut.PresetTriggerCmd, M1_PresetValueOut := encoderM1.HwOut.PresetValueOut, M2_PresetTriggerCmd := encoderM2.HwOut.PresetTriggerCmd, M2_PresetValueOut := encoderM2.HwOut.PresetValueOut, RawPosM1 := raw1, RawPosM2 := raw2); raw1 := bench.RawPosM1; raw2 := bench.RawPosM2;
hw1.RawPosIn := bench.Winch.COD1_PosValue; hw1.SlaveOperational := TRUE; hw2.RawPosIn := bench.Winch.COD2_PosValue; hw2.SlaveOperational := TRUE;
encoderM1(Enable := TRUE, HomingPermit := TRUE, HomingAtTargetM := btnM1, CfgHomingTargetM := 8.7, CfgTopSensorPosM := 8.7, HwIn := hw1, Cfg := cfgEncoder, Calib := calibM1); calibM1 := encoderM1.Calib;
bucketEdge(CLK := btnBucket);
encoderM2(Enable := TRUE, HomingPermit := TRUE, HomingAtTargetM := btnM2 OR bucketEdge.Q, CfgHomingTargetM := 23.7, CfgTopSensorPosM := 23.7, UseDynamicTarget := bucketEdge.Q, DynamicHomingTargetM := encoderM1.Measurement.CablePosM + cfgBucket.OffsetCloseM, HwIn := hw2, Cfg := cfgEncoder, Calib := calibM2); calibM2 := encoderM2.Calib;
bucket(Enable := TRUE, Mode := E_Mode.MAINT_N2, PowerContactorEngaged := TRUE, CablePosM1 := encoderM1.Measurement.CablePosM, CablePosM2 := encoderM2.Measurement.CablePosM, HomedM1 := encoderM1.Homed, HomedM2 := encoderM2.Homed, HomedAndReliableM1 := encoderM1.HomedAndReliable, HomedAndReliableM2 := encoderM2.HomedAndReliable, HomingSuspectM1 := encoderM1.HomingSuspect, HomingSuspectM2 := encoderM2.HomingSuspect, ConfirmClosePosition := btnBucket, Config := cfgBucket, BucketState := bucketState); bucketState := bucket.BucketState;
home.M1Status.HomedAndReliable := encoderM1.HomedAndReliable; home.M2Status.HomedAndReliable := encoderM2.HomedAndReliable; home(BucketOffsetValid := bucketState.BucketReferenced, BtnValidation := bench.Operator.JoyBtnRaw);
ADVANCE_TIME(10000000);
bench(M1_PresetTriggerCmd := encoderM1.HwOut.PresetTriggerCmd, M1_PresetValueOut := encoderM1.HwOut.PresetValueOut, M2_PresetTriggerCmd := encoderM2.HwOut.PresetTriggerCmd, M2_PresetValueOut := encoderM2.HwOut.PresetValueOut, RawPosM1 := raw1, RawPosM2 := raw2); raw1 := bench.RawPosM1; raw2 := bench.RawPosM2;
hw1.RawPosIn := bench.Winch.COD1_PosValue; hw1.SlaveOperational := TRUE; hw2.RawPosIn := bench.Winch.COD2_PosValue; hw2.SlaveOperational := TRUE;
encoderM1(Enable := TRUE, HomingPermit := TRUE, HomingAtTargetM := btnM1, CfgHomingTargetM := 8.7, CfgTopSensorPosM := 8.7, HwIn := hw1, Cfg := cfgEncoder, Calib := calibM1); calibM1 := encoderM1.Calib;
bucketEdge(CLK := btnBucket);
encoderM2(Enable := TRUE, HomingPermit := TRUE, HomingAtTargetM := btnM2 OR bucketEdge.Q, CfgHomingTargetM := 23.7, CfgTopSensorPosM := 23.7, UseDynamicTarget := bucketEdge.Q, DynamicHomingTargetM := encoderM1.Measurement.CablePosM + cfgBucket.OffsetCloseM, HwIn := hw2, Cfg := cfgEncoder, Calib := calibM2); calibM2 := encoderM2.Calib;
bucket(Enable := TRUE, Mode := E_Mode.MAINT_N2, PowerContactorEngaged := TRUE, CablePosM1 := encoderM1.Measurement.CablePosM, CablePosM2 := encoderM2.Measurement.CablePosM, HomedM1 := encoderM1.Homed, HomedM2 := encoderM2.Homed, HomedAndReliableM1 := encoderM1.HomedAndReliable, HomedAndReliableM2 := encoderM2.HomedAndReliable, HomingSuspectM1 := encoderM1.HomingSuspect, HomingSuspectM2 := encoderM2.HomingSuspect, ConfirmClosePosition := btnBucket, Config := cfgBucket, BucketState := bucketState); bucketState := bucket.BucketState;
home.M1Status.HomedAndReliable := encoderM1.HomedAndReliable; home.M2Status.HomedAndReliable := encoderM2.HomedAndReliable; home(BucketOffsetValid := bucketState.BucketReferenced, BtnValidation := bench.Operator.JoyBtnRaw);
ADVANCE_TIME(10000000);
bench(M1_PresetTriggerCmd := encoderM1.HwOut.PresetTriggerCmd, M1_PresetValueOut := encoderM1.HwOut.PresetValueOut, M2_PresetTriggerCmd := encoderM2.HwOut.PresetTriggerCmd, M2_PresetValueOut := encoderM2.HwOut.PresetValueOut, RawPosM1 := raw1, RawPosM2 := raw2); raw1 := bench.RawPosM1; raw2 := bench.RawPosM2;
hw1.RawPosIn := bench.Winch.COD1_PosValue; hw1.SlaveOperational := TRUE; hw2.RawPosIn := bench.Winch.COD2_PosValue; hw2.SlaveOperational := TRUE;
encoderM1(Enable := TRUE, HomingPermit := TRUE, HomingAtTargetM := btnM1, CfgHomingTargetM := 8.7, CfgTopSensorPosM := 8.7, HwIn := hw1, Cfg := cfgEncoder, Calib := calibM1); calibM1 := encoderM1.Calib;
bucketEdge(CLK := btnBucket);
encoderM2(Enable := TRUE, HomingPermit := TRUE, HomingAtTargetM := btnM2 OR bucketEdge.Q, CfgHomingTargetM := 23.7, CfgTopSensorPosM := 23.7, UseDynamicTarget := bucketEdge.Q, DynamicHomingTargetM := encoderM1.Measurement.CablePosM + cfgBucket.OffsetCloseM, HwIn := hw2, Cfg := cfgEncoder, Calib := calibM2); calibM2 := encoderM2.Calib;
bucket(Enable := TRUE, Mode := E_Mode.MAINT_N2, PowerContactorEngaged := TRUE, CablePosM1 := encoderM1.Measurement.CablePosM, CablePosM2 := encoderM2.Measurement.CablePosM, HomedM1 := encoderM1.Homed, HomedM2 := encoderM2.Homed, HomedAndReliableM1 := encoderM1.HomedAndReliable, HomedAndReliableM2 := encoderM2.HomedAndReliable, HomingSuspectM1 := encoderM1.HomingSuspect, HomingSuspectM2 := encoderM2.HomingSuspect, ConfirmClosePosition := btnBucket, Config := cfgBucket, BucketState := bucketState); bucketState := bucket.BucketState;
home.M1Status.HomedAndReliable := encoderM1.HomedAndReliable; home.M2Status.HomedAndReliable := encoderM2.HomedAndReliable; home(BucketOffsetValid := bucketState.BucketReferenced, BtnValidation := bench.Operator.JoyBtnRaw);
ADVANCE_TIME(10000000);
bench(M1_PresetTriggerCmd := encoderM1.HwOut.PresetTriggerCmd, M1_PresetValueOut := encoderM1.HwOut.PresetValueOut, M2_PresetTriggerCmd := encoderM2.HwOut.PresetTriggerCmd, M2_PresetValueOut := encoderM2.HwOut.PresetValueOut, RawPosM1 := raw1, RawPosM2 := raw2); raw1 := bench.RawPosM1; raw2 := bench.RawPosM2;
hw1.RawPosIn := bench.Winch.COD1_PosValue; hw1.SlaveOperational := TRUE; hw2.RawPosIn := bench.Winch.COD2_PosValue; hw2.SlaveOperational := TRUE;
encoderM1(Enable := TRUE, HomingPermit := TRUE, HomingAtTargetM := btnM1, CfgHomingTargetM := 8.7, CfgTopSensorPosM := 8.7, HwIn := hw1, Cfg := cfgEncoder, Calib := calibM1); calibM1 := encoderM1.Calib;
bucketEdge(CLK := btnBucket);
encoderM2(Enable := TRUE, HomingPermit := TRUE, HomingAtTargetM := btnM2 OR bucketEdge.Q, CfgHomingTargetM := 23.7, CfgTopSensorPosM := 23.7, UseDynamicTarget := bucketEdge.Q, DynamicHomingTargetM := encoderM1.Measurement.CablePosM + cfgBucket.OffsetCloseM, HwIn := hw2, Cfg := cfgEncoder, Calib := calibM2); calibM2 := encoderM2.Calib;
bucket(Enable := TRUE, Mode := E_Mode.MAINT_N2, PowerContactorEngaged := TRUE, CablePosM1 := encoderM1.Measurement.CablePosM, CablePosM2 := encoderM2.Measurement.CablePosM, HomedM1 := encoderM1.Homed, HomedM2 := encoderM2.Homed, HomedAndReliableM1 := encoderM1.HomedAndReliable, HomedAndReliableM2 := encoderM2.HomedAndReliable, HomingSuspectM1 := encoderM1.HomingSuspect, HomingSuspectM2 := encoderM2.HomingSuspect, ConfirmClosePosition := btnBucket, Config := cfgBucket, BucketState := bucketState); bucketState := bucket.BucketState;
home.M1Status.HomedAndReliable := encoderM1.HomedAndReliable; home.M2Status.HomedAndReliable := encoderM2.HomedAndReliable; home(BucketOffsetValid := bucketState.BucketReferenced, BtnValidation := bench.Operator.JoyBtnRaw);
ADVANCE_TIME(10000000);
bench(M1_PresetTriggerCmd := encoderM1.HwOut.PresetTriggerCmd, M1_PresetValueOut := encoderM1.HwOut.PresetValueOut, M2_PresetTriggerCmd := encoderM2.HwOut.PresetTriggerCmd, M2_PresetValueOut := encoderM2.HwOut.PresetValueOut, RawPosM1 := raw1, RawPosM2 := raw2); raw1 := bench.RawPosM1; raw2 := bench.RawPosM2;
hw1.RawPosIn := bench.Winch.COD1_PosValue; hw1.SlaveOperational := TRUE; hw2.RawPosIn := bench.Winch.COD2_PosValue; hw2.SlaveOperational := TRUE;
encoderM1(Enable := TRUE, HomingPermit := TRUE, HomingAtTargetM := btnM1, CfgHomingTargetM := 8.7, CfgTopSensorPosM := 8.7, HwIn := hw1, Cfg := cfgEncoder, Calib := calibM1); calibM1 := encoderM1.Calib;
bucketEdge(CLK := btnBucket);
encoderM2(Enable := TRUE, HomingPermit := TRUE, HomingAtTargetM := btnM2 OR bucketEdge.Q, CfgHomingTargetM := 23.7, CfgTopSensorPosM := 23.7, UseDynamicTarget := bucketEdge.Q, DynamicHomingTargetM := encoderM1.Measurement.CablePosM + cfgBucket.OffsetCloseM, HwIn := hw2, Cfg := cfgEncoder, Calib := calibM2); calibM2 := encoderM2.Calib;
bucket(Enable := TRUE, Mode := E_Mode.MAINT_N2, PowerContactorEngaged := TRUE, CablePosM1 := encoderM1.Measurement.CablePosM, CablePosM2 := encoderM2.Measurement.CablePosM, HomedM1 := encoderM1.Homed, HomedM2 := encoderM2.Homed, HomedAndReliableM1 := encoderM1.HomedAndReliable, HomedAndReliableM2 := encoderM2.HomedAndReliable, HomingSuspectM1 := encoderM1.HomingSuspect, HomingSuspectM2 := encoderM2.HomingSuspect, ConfirmClosePosition := btnBucket, Config := cfgBucket, BucketState := bucketState); bucketState := bucket.BucketState;
home.M1Status.HomedAndReliable := encoderM1.HomedAndReliable; home.M2Status.HomedAndReliable := encoderM2.HomedAndReliable; home(BucketOffsetValid := bucketState.BucketReferenced, BtnValidation := bench.Operator.JoyBtnRaw);
ADVANCE_TIME(10000000);
bench(M1_PresetTriggerCmd := encoderM1.HwOut.PresetTriggerCmd, M1_PresetValueOut := encoderM1.HwOut.PresetValueOut, M2_PresetTriggerCmd := encoderM2.HwOut.PresetTriggerCmd, M2_PresetValueOut := encoderM2.HwOut.PresetValueOut, RawPosM1 := raw1, RawPosM2 := raw2); raw1 := bench.RawPosM1; raw2 := bench.RawPosM2;
hw1.RawPosIn := bench.Winch.COD1_PosValue; hw1.SlaveOperational := TRUE; hw2.RawPosIn := bench.Winch.COD2_PosValue; hw2.SlaveOperational := TRUE;
encoderM1(Enable := TRUE, HomingPermit := TRUE, HomingAtTargetM := btnM1, CfgHomingTargetM := 8.7, CfgTopSensorPosM := 8.7, HwIn := hw1, Cfg := cfgEncoder, Calib := calibM1); calibM1 := encoderM1.Calib;
bucketEdge(CLK := btnBucket);
encoderM2(Enable := TRUE, HomingPermit := TRUE, HomingAtTargetM := btnM2 OR bucketEdge.Q, CfgHomingTargetM := 23.7, CfgTopSensorPosM := 23.7, UseDynamicTarget := bucketEdge.Q, DynamicHomingTargetM := encoderM1.Measurement.CablePosM + cfgBucket.OffsetCloseM, HwIn := hw2, Cfg := cfgEncoder, Calib := calibM2); calibM2 := encoderM2.Calib;
bucket(Enable := TRUE, Mode := E_Mode.MAINT_N2, PowerContactorEngaged := TRUE, CablePosM1 := encoderM1.Measurement.CablePosM, CablePosM2 := encoderM2.Measurement.CablePosM, HomedM1 := encoderM1.Homed, HomedM2 := encoderM2.Homed, HomedAndReliableM1 := encoderM1.HomedAndReliable, HomedAndReliableM2 := encoderM2.HomedAndReliable, HomingSuspectM1 := encoderM1.HomingSuspect, HomingSuspectM2 := encoderM2.HomingSuspect, ConfirmClosePosition := btnBucket, Config := cfgBucket, BucketState := bucketState); bucketState := bucket.BucketState;
home.M1Status.HomedAndReliable := encoderM1.HomedAndReliable; home.M2Status.HomedAndReliable := encoderM2.HomedAndReliable; home(BucketOffsetValid := bucketState.BucketReferenced, BtnValidation := bench.Operator.JoyBtnRaw);
ADVANCE_TIME(10000000);
bench(M1_PresetTriggerCmd := encoderM1.HwOut.PresetTriggerCmd, M1_PresetValueOut := encoderM1.HwOut.PresetValueOut, M2_PresetTriggerCmd := encoderM2.HwOut.PresetTriggerCmd, M2_PresetValueOut := encoderM2.HwOut.PresetValueOut, RawPosM1 := raw1, RawPosM2 := raw2); raw1 := bench.RawPosM1; raw2 := bench.RawPosM2;
hw1.RawPosIn := bench.Winch.COD1_PosValue; hw1.SlaveOperational := TRUE; hw2.RawPosIn := bench.Winch.COD2_PosValue; hw2.SlaveOperational := TRUE;
encoderM1(Enable := TRUE, HomingPermit := TRUE, HomingAtTargetM := btnM1, CfgHomingTargetM := 8.7, CfgTopSensorPosM := 8.7, HwIn := hw1, Cfg := cfgEncoder, Calib := calibM1); calibM1 := encoderM1.Calib;
bucketEdge(CLK := btnBucket);
encoderM2(Enable := TRUE, HomingPermit := TRUE, HomingAtTargetM := btnM2 OR bucketEdge.Q, CfgHomingTargetM := 23.7, CfgTopSensorPosM := 23.7, UseDynamicTarget := bucketEdge.Q, DynamicHomingTargetM := encoderM1.Measurement.CablePosM + cfgBucket.OffsetCloseM, HwIn := hw2, Cfg := cfgEncoder, Calib := calibM2); calibM2 := encoderM2.Calib;
bucket(Enable := TRUE, Mode := E_Mode.MAINT_N2, PowerContactorEngaged := TRUE, CablePosM1 := encoderM1.Measurement.CablePosM, CablePosM2 := encoderM2.Measurement.CablePosM, HomedM1 := encoderM1.Homed, HomedM2 := encoderM2.Homed, HomedAndReliableM1 := encoderM1.HomedAndReliable, HomedAndReliableM2 := encoderM2.HomedAndReliable, HomingSuspectM1 := encoderM1.HomingSuspect, HomingSuspectM2 := encoderM2.HomingSuspect, ConfirmClosePosition := btnBucket, Config := cfgBucket, BucketState := bucketState); bucketState := bucket.BucketState;
home.M1Status.HomedAndReliable := encoderM1.HomedAndReliable; home.M2Status.HomedAndReliable := encoderM2.HomedAndReliable; home(BucketOffsetValid := bucketState.BucketReferenced, BtnValidation := bench.Operator.JoyBtnRaw);
ADVANCE_TIME(10000000);
bench(M1_PresetTriggerCmd := encoderM1.HwOut.PresetTriggerCmd, M1_PresetValueOut := encoderM1.HwOut.PresetValueOut, M2_PresetTriggerCmd := encoderM2.HwOut.PresetTriggerCmd, M2_PresetValueOut := encoderM2.HwOut.PresetValueOut, RawPosM1 := raw1, RawPosM2 := raw2); raw1 := bench.RawPosM1; raw2 := bench.RawPosM2;
hw1.RawPosIn := bench.Winch.COD1_PosValue; hw1.SlaveOperational := TRUE; hw2.RawPosIn := bench.Winch.COD2_PosValue; hw2.SlaveOperational := TRUE;
encoderM1(Enable := TRUE, HomingPermit := TRUE, HomingAtTargetM := btnM1, CfgHomingTargetM := 8.7, CfgTopSensorPosM := 8.7, HwIn := hw1, Cfg := cfgEncoder, Calib := calibM1); calibM1 := encoderM1.Calib;
bucketEdge(CLK := btnBucket);
encoderM2(Enable := TRUE, HomingPermit := TRUE, HomingAtTargetM := btnM2 OR bucketEdge.Q, CfgHomingTargetM := 23.7, CfgTopSensorPosM := 23.7, UseDynamicTarget := bucketEdge.Q, DynamicHomingTargetM := encoderM1.Measurement.CablePosM + cfgBucket.OffsetCloseM, HwIn := hw2, Cfg := cfgEncoder, Calib := calibM2); calibM2 := encoderM2.Calib;
bucket(Enable := TRUE, Mode := E_Mode.MAINT_N2, PowerContactorEngaged := TRUE, CablePosM1 := encoderM1.Measurement.CablePosM, CablePosM2 := encoderM2.Measurement.CablePosM, HomedM1 := encoderM1.Homed, HomedM2 := encoderM2.Homed, HomedAndReliableM1 := encoderM1.HomedAndReliable, HomedAndReliableM2 := encoderM2.HomedAndReliable, HomingSuspectM1 := encoderM1.HomingSuspect, HomingSuspectM2 := encoderM2.HomingSuspect, ConfirmClosePosition := btnBucket, Config := cfgBucket, BucketState := bucketState); bucketState := bucket.BucketState;
home.M1Status.HomedAndReliable := encoderM1.HomedAndReliable; home.M2Status.HomedAndReliable := encoderM2.HomedAndReliable; home(BucketOffsetValid := bucketState.BucketReferenced, BtnValidation := bench.Operator.JoyBtnRaw);
ADVANCE_TIME(10000000);
bench(M1_PresetTriggerCmd := encoderM1.HwOut.PresetTriggerCmd, M1_PresetValueOut := encoderM1.HwOut.PresetValueOut, M2_PresetTriggerCmd := encoderM2.HwOut.PresetTriggerCmd, M2_PresetValueOut := encoderM2.HwOut.PresetValueOut, RawPosM1 := raw1, RawPosM2 := raw2); raw1 := bench.RawPosM1; raw2 := bench.RawPosM2;
hw1.RawPosIn := bench.Winch.COD1_PosValue; hw1.SlaveOperational := TRUE; hw2.RawPosIn := bench.Winch.COD2_PosValue; hw2.SlaveOperational := TRUE;
encoderM1(Enable := TRUE, HomingPermit := TRUE, HomingAtTargetM := btnM1, CfgHomingTargetM := 8.7, CfgTopSensorPosM := 8.7, HwIn := hw1, Cfg := cfgEncoder, Calib := calibM1); calibM1 := encoderM1.Calib;
bucketEdge(CLK := btnBucket);
encoderM2(Enable := TRUE, HomingPermit := TRUE, HomingAtTargetM := btnM2 OR bucketEdge.Q, CfgHomingTargetM := 23.7, CfgTopSensorPosM := 23.7, UseDynamicTarget := bucketEdge.Q, DynamicHomingTargetM := encoderM1.Measurement.CablePosM + cfgBucket.OffsetCloseM, HwIn := hw2, Cfg := cfgEncoder, Calib := calibM2); calibM2 := encoderM2.Calib;
bucket(Enable := TRUE, Mode := E_Mode.MAINT_N2, PowerContactorEngaged := TRUE, CablePosM1 := encoderM1.Measurement.CablePosM, CablePosM2 := encoderM2.Measurement.CablePosM, HomedM1 := encoderM1.Homed, HomedM2 := encoderM2.Homed, HomedAndReliableM1 := encoderM1.HomedAndReliable, HomedAndReliableM2 := encoderM2.HomedAndReliable, HomingSuspectM1 := encoderM1.HomingSuspect, HomingSuspectM2 := encoderM2.HomingSuspect, ConfirmClosePosition := btnBucket, Config := cfgBucket, BucketState := bucketState); bucketState := bucket.BucketState;
home.M1Status.HomedAndReliable := encoderM1.HomedAndReliable; home.M2Status.HomedAndReliable := encoderM2.HomedAndReliable; home(BucketOffsetValid := bucketState.BucketReferenced, BtnValidation := bench.Operator.JoyBtnRaw);
ADVANCE_TIME(10000000);
bench(M1_PresetTriggerCmd := encoderM1.HwOut.PresetTriggerCmd, M1_PresetValueOut := encoderM1.HwOut.PresetValueOut, M2_PresetTriggerCmd := encoderM2.HwOut.PresetTriggerCmd, M2_PresetValueOut := encoderM2.HwOut.PresetValueOut, RawPosM1 := raw1, RawPosM2 := raw2); raw1 := bench.RawPosM1; raw2 := bench.RawPosM2;
hw1.RawPosIn := bench.Winch.COD1_PosValue; hw1.SlaveOperational := TRUE; hw2.RawPosIn := bench.Winch.COD2_PosValue; hw2.SlaveOperational := TRUE;
encoderM1(Enable := TRUE, HomingPermit := TRUE, HomingAtTargetM := btnM1, CfgHomingTargetM := 8.7, CfgTopSensorPosM := 8.7, HwIn := hw1, Cfg := cfgEncoder, Calib := calibM1); calibM1 := encoderM1.Calib;
bucketEdge(CLK := btnBucket);
encoderM2(Enable := TRUE, HomingPermit := TRUE, HomingAtTargetM := btnM2 OR bucketEdge.Q, CfgHomingTargetM := 23.7, CfgTopSensorPosM := 23.7, UseDynamicTarget := bucketEdge.Q, DynamicHomingTargetM := encoderM1.Measurement.CablePosM + cfgBucket.OffsetCloseM, HwIn := hw2, Cfg := cfgEncoder, Calib := calibM2); calibM2 := encoderM2.Calib;
bucket(Enable := TRUE, Mode := E_Mode.MAINT_N2, PowerContactorEngaged := TRUE, CablePosM1 := encoderM1.Measurement.CablePosM, CablePosM2 := encoderM2.Measurement.CablePosM, HomedM1 := encoderM1.Homed, HomedM2 := encoderM2.Homed, HomedAndReliableM1 := encoderM1.HomedAndReliable, HomedAndReliableM2 := encoderM2.HomedAndReliable, HomingSuspectM1 := encoderM1.HomingSuspect, HomingSuspectM2 := encoderM2.HomingSuspect, ConfirmClosePosition := btnBucket, Config := cfgBucket, BucketState := bucketState); bucketState := bucket.BucketState;
home.M1Status.HomedAndReliable := encoderM1.HomedAndReliable; home.M2Status.HomedAndReliable := encoderM2.HomedAndReliable; home(BucketOffsetValid := bucketState.BucketReferenced, BtnValidation := bench.Operator.JoyBtnRaw);
ADVANCE_TIME(10000000);
bench(M1_PresetTriggerCmd := encoderM1.HwOut.PresetTriggerCmd, M1_PresetValueOut := encoderM1.HwOut.PresetValueOut, M2_PresetTriggerCmd := encoderM2.HwOut.PresetTriggerCmd, M2_PresetValueOut := encoderM2.HwOut.PresetValueOut, RawPosM1 := raw1, RawPosM2 := raw2); raw1 := bench.RawPosM1; raw2 := bench.RawPosM2;
hw1.RawPosIn := bench.Winch.COD1_PosValue; hw1.SlaveOperational := TRUE; hw2.RawPosIn := bench.Winch.COD2_PosValue; hw2.SlaveOperational := TRUE;
encoderM1(Enable := TRUE, HomingPermit := TRUE, HomingAtTargetM := btnM1, CfgHomingTargetM := 8.7, CfgTopSensorPosM := 8.7, HwIn := hw1, Cfg := cfgEncoder, Calib := calibM1); calibM1 := encoderM1.Calib;
bucketEdge(CLK := btnBucket);
encoderM2(Enable := TRUE, HomingPermit := TRUE, HomingAtTargetM := btnM2 OR bucketEdge.Q, CfgHomingTargetM := 23.7, CfgTopSensorPosM := 23.7, UseDynamicTarget := bucketEdge.Q, DynamicHomingTargetM := encoderM1.Measurement.CablePosM + cfgBucket.OffsetCloseM, HwIn := hw2, Cfg := cfgEncoder, Calib := calibM2); calibM2 := encoderM2.Calib;
bucket(Enable := TRUE, Mode := E_Mode.MAINT_N2, PowerContactorEngaged := TRUE, CablePosM1 := encoderM1.Measurement.CablePosM, CablePosM2 := encoderM2.Measurement.CablePosM, HomedM1 := encoderM1.Homed, HomedM2 := encoderM2.Homed, HomedAndReliableM1 := encoderM1.HomedAndReliable, HomedAndReliableM2 := encoderM2.HomedAndReliable, HomingSuspectM1 := encoderM1.HomingSuspect, HomingSuspectM2 := encoderM2.HomingSuspect, ConfirmClosePosition := btnBucket, Config := cfgBucket, BucketState := bucketState); bucketState := bucket.BucketState;
home.M1Status.HomedAndReliable := encoderM1.HomedAndReliable; home.M2Status.HomedAndReliable := encoderM2.HomedAndReliable; home(BucketOffsetValid := bucketState.BucketReferenced, BtnValidation := bench.Operator.JoyBtnRaw);
ADVANCE_TIME(10000000);
bench(M1_PresetTriggerCmd := encoderM1.HwOut.PresetTriggerCmd, M1_PresetValueOut := encoderM1.HwOut.PresetValueOut, M2_PresetTriggerCmd := encoderM2.HwOut.PresetTriggerCmd, M2_PresetValueOut := encoderM2.HwOut.PresetValueOut, RawPosM1 := raw1, RawPosM2 := raw2); raw1 := bench.RawPosM1; raw2 := bench.RawPosM2;
hw1.RawPosIn := bench.Winch.COD1_PosValue; hw1.SlaveOperational := TRUE; hw2.RawPosIn := bench.Winch.COD2_PosValue; hw2.SlaveOperational := TRUE;
encoderM1(Enable := TRUE, HomingPermit := TRUE, HomingAtTargetM := btnM1, CfgHomingTargetM := 8.7, CfgTopSensorPosM := 8.7, HwIn := hw1, Cfg := cfgEncoder, Calib := calibM1); calibM1 := encoderM1.Calib;
bucketEdge(CLK := btnBucket);
encoderM2(Enable := TRUE, HomingPermit := TRUE, HomingAtTargetM := btnM2 OR bucketEdge.Q, CfgHomingTargetM := 23.7, CfgTopSensorPosM := 23.7, UseDynamicTarget := bucketEdge.Q, DynamicHomingTargetM := encoderM1.Measurement.CablePosM + cfgBucket.OffsetCloseM, HwIn := hw2, Cfg := cfgEncoder, Calib := calibM2); calibM2 := encoderM2.Calib;
bucket(Enable := TRUE, Mode := E_Mode.MAINT_N2, PowerContactorEngaged := TRUE, CablePosM1 := encoderM1.Measurement.CablePosM, CablePosM2 := encoderM2.Measurement.CablePosM, HomedM1 := encoderM1.Homed, HomedM2 := encoderM2.Homed, HomedAndReliableM1 := encoderM1.HomedAndReliable, HomedAndReliableM2 := encoderM2.HomedAndReliable, HomingSuspectM1 := encoderM1.HomingSuspect, HomingSuspectM2 := encoderM2.HomingSuspect, ConfirmClosePosition := btnBucket, Config := cfgBucket, BucketState := bucketState); bucketState := bucket.BucketState;
home.M1Status.HomedAndReliable := encoderM1.HomedAndReliable; home.M2Status.HomedAndReliable := encoderM2.HomedAndReliable; home(BucketOffsetValid := bucketState.BucketReferenced, BtnValidation := bench.Operator.JoyBtnRaw);
ADVANCE_TIME(10000000);
bench(M1_PresetTriggerCmd := encoderM1.HwOut.PresetTriggerCmd, M1_PresetValueOut := encoderM1.HwOut.PresetValueOut, M2_PresetTriggerCmd := encoderM2.HwOut.PresetTriggerCmd, M2_PresetValueOut := encoderM2.HwOut.PresetValueOut, RawPosM1 := raw1, RawPosM2 := raw2); raw1 := bench.RawPosM1; raw2 := bench.RawPosM2;
hw1.RawPosIn := bench.Winch.COD1_PosValue; hw1.SlaveOperational := TRUE; hw2.RawPosIn := bench.Winch.COD2_PosValue; hw2.SlaveOperational := TRUE;
encoderM1(Enable := TRUE, HomingPermit := TRUE, HomingAtTargetM := btnM1, CfgHomingTargetM := 8.7, CfgTopSensorPosM := 8.7, HwIn := hw1, Cfg := cfgEncoder, Calib := calibM1); calibM1 := encoderM1.Calib;
bucketEdge(CLK := btnBucket);
encoderM2(Enable := TRUE, HomingPermit := TRUE, HomingAtTargetM := btnM2 OR bucketEdge.Q, CfgHomingTargetM := 23.7, CfgTopSensorPosM := 23.7, UseDynamicTarget := bucketEdge.Q, DynamicHomingTargetM := encoderM1.Measurement.CablePosM + cfgBucket.OffsetCloseM, HwIn := hw2, Cfg := cfgEncoder, Calib := calibM2); calibM2 := encoderM2.Calib;
bucket(Enable := TRUE, Mode := E_Mode.MAINT_N2, PowerContactorEngaged := TRUE, CablePosM1 := encoderM1.Measurement.CablePosM, CablePosM2 := encoderM2.Measurement.CablePosM, HomedM1 := encoderM1.Homed, HomedM2 := encoderM2.Homed, HomedAndReliableM1 := encoderM1.HomedAndReliable, HomedAndReliableM2 := encoderM2.HomedAndReliable, HomingSuspectM1 := encoderM1.HomingSuspect, HomingSuspectM2 := encoderM2.HomingSuspect, ConfirmClosePosition := btnBucket, Config := cfgBucket, BucketState := bucketState); bucketState := bucket.BucketState;
home.M1Status.HomedAndReliable := encoderM1.HomedAndReliable; home.M2Status.HomedAndReliable := encoderM2.HomedAndReliable; home(BucketOffsetValid := bucketState.BucketReferenced, BtnValidation := bench.Operator.JoyBtnRaw);
ADVANCE_TIME(10000000);
bench(M1_PresetTriggerCmd := encoderM1.HwOut.PresetTriggerCmd, M1_PresetValueOut := encoderM1.HwOut.PresetValueOut, M2_PresetTriggerCmd := encoderM2.HwOut.PresetTriggerCmd, M2_PresetValueOut := encoderM2.HwOut.PresetValueOut, RawPosM1 := raw1, RawPosM2 := raw2); raw1 := bench.RawPosM1; raw2 := bench.RawPosM2;
hw1.RawPosIn := bench.Winch.COD1_PosValue; hw1.SlaveOperational := TRUE; hw2.RawPosIn := bench.Winch.COD2_PosValue; hw2.SlaveOperational := TRUE;
encoderM1(Enable := TRUE, HomingPermit := TRUE, HomingAtTargetM := btnM1, CfgHomingTargetM := 8.7, CfgTopSensorPosM := 8.7, HwIn := hw1, Cfg := cfgEncoder, Calib := calibM1); calibM1 := encoderM1.Calib;
bucketEdge(CLK := btnBucket);
encoderM2(Enable := TRUE, HomingPermit := TRUE, HomingAtTargetM := btnM2 OR bucketEdge.Q, CfgHomingTargetM := 23.7, CfgTopSensorPosM := 23.7, UseDynamicTarget := bucketEdge.Q, DynamicHomingTargetM := encoderM1.Measurement.CablePosM + cfgBucket.OffsetCloseM, HwIn := hw2, Cfg := cfgEncoder, Calib := calibM2); calibM2 := encoderM2.Calib;
bucket(Enable := TRUE, Mode := E_Mode.MAINT_N2, PowerContactorEngaged := TRUE, CablePosM1 := encoderM1.Measurement.CablePosM, CablePosM2 := encoderM2.Measurement.CablePosM, HomedM1 := encoderM1.Homed, HomedM2 := encoderM2.Homed, HomedAndReliableM1 := encoderM1.HomedAndReliable, HomedAndReliableM2 := encoderM2.HomedAndReliable, HomingSuspectM1 := encoderM1.HomingSuspect, HomingSuspectM2 := encoderM2.HomingSuspect, ConfirmClosePosition := btnBucket, Config := cfgBucket, BucketState := bucketState); bucketState := bucket.BucketState;
home.M1Status.HomedAndReliable := encoderM1.HomedAndReliable; home.M2Status.HomedAndReliable := encoderM2.HomedAndReliable; home(BucketOffsetValid := bucketState.BucketReferenced, BtnValidation := bench.Operator.JoyBtnRaw);
ADVANCE_TIME(10000000);
bench(M1_PresetTriggerCmd := encoderM1.HwOut.PresetTriggerCmd, M1_PresetValueOut := encoderM1.HwOut.PresetValueOut, M2_PresetTriggerCmd := encoderM2.HwOut.PresetTriggerCmd, M2_PresetValueOut := encoderM2.HwOut.PresetValueOut, RawPosM1 := raw1, RawPosM2 := raw2); raw1 := bench.RawPosM1; raw2 := bench.RawPosM2;
hw1.RawPosIn := bench.Winch.COD1_PosValue; hw1.SlaveOperational := TRUE; hw2.RawPosIn := bench.Winch.COD2_PosValue; hw2.SlaveOperational := TRUE;
encoderM1(Enable := TRUE, HomingPermit := TRUE, HomingAtTargetM := btnM1, CfgHomingTargetM := 8.7, CfgTopSensorPosM := 8.7, HwIn := hw1, Cfg := cfgEncoder, Calib := calibM1); calibM1 := encoderM1.Calib;
bucketEdge(CLK := btnBucket);
encoderM2(Enable := TRUE, HomingPermit := TRUE, HomingAtTargetM := btnM2 OR bucketEdge.Q, CfgHomingTargetM := 23.7, CfgTopSensorPosM := 23.7, UseDynamicTarget := bucketEdge.Q, DynamicHomingTargetM := encoderM1.Measurement.CablePosM + cfgBucket.OffsetCloseM, HwIn := hw2, Cfg := cfgEncoder, Calib := calibM2); calibM2 := encoderM2.Calib;
bucket(Enable := TRUE, Mode := E_Mode.MAINT_N2, PowerContactorEngaged := TRUE, CablePosM1 := encoderM1.Measurement.CablePosM, CablePosM2 := encoderM2.Measurement.CablePosM, HomedM1 := encoderM1.Homed, HomedM2 := encoderM2.Homed, HomedAndReliableM1 := encoderM1.HomedAndReliable, HomedAndReliableM2 := encoderM2.HomedAndReliable, HomingSuspectM1 := encoderM1.HomingSuspect, HomingSuspectM2 := encoderM2.HomingSuspect, ConfirmClosePosition := btnBucket, Config := cfgBucket, BucketState := bucketState); bucketState := bucket.BucketState;
home.M1Status.HomedAndReliable := encoderM1.HomedAndReliable; home.M2Status.HomedAndReliable := encoderM2.HomedAndReliable; home(BucketOffsetValid := bucketState.BucketReferenced, BtnValidation := bench.Operator.JoyBtnRaw);
ADVANCE_TIME(10000000);
bench(M1_PresetTriggerCmd := encoderM1.HwOut.PresetTriggerCmd, M1_PresetValueOut := encoderM1.HwOut.PresetValueOut, M2_PresetTriggerCmd := encoderM2.HwOut.PresetTriggerCmd, M2_PresetValueOut := encoderM2.HwOut.PresetValueOut, RawPosM1 := raw1, RawPosM2 := raw2); raw1 := bench.RawPosM1; raw2 := bench.RawPosM2;
hw1.RawPosIn := bench.Winch.COD1_PosValue; hw1.SlaveOperational := TRUE; hw2.RawPosIn := bench.Winch.COD2_PosValue; hw2.SlaveOperational := TRUE;
encoderM1(Enable := TRUE, HomingPermit := TRUE, HomingAtTargetM := btnM1, CfgHomingTargetM := 8.7, CfgTopSensorPosM := 8.7, HwIn := hw1, Cfg := cfgEncoder, Calib := calibM1); calibM1 := encoderM1.Calib;
bucketEdge(CLK := btnBucket);
encoderM2(Enable := TRUE, HomingPermit := TRUE, HomingAtTargetM := btnM2 OR bucketEdge.Q, CfgHomingTargetM := 23.7, CfgTopSensorPosM := 23.7, UseDynamicTarget := bucketEdge.Q, DynamicHomingTargetM := encoderM1.Measurement.CablePosM + cfgBucket.OffsetCloseM, HwIn := hw2, Cfg := cfgEncoder, Calib := calibM2); calibM2 := encoderM2.Calib;
bucket(Enable := TRUE, Mode := E_Mode.MAINT_N2, PowerContactorEngaged := TRUE, CablePosM1 := encoderM1.Measurement.CablePosM, CablePosM2 := encoderM2.Measurement.CablePosM, HomedM1 := encoderM1.Homed, HomedM2 := encoderM2.Homed, HomedAndReliableM1 := encoderM1.HomedAndReliable, HomedAndReliableM2 := encoderM2.HomedAndReliable, HomingSuspectM1 := encoderM1.HomingSuspect, HomingSuspectM2 := encoderM2.HomingSuspect, ConfirmClosePosition := btnBucket, Config := cfgBucket, BucketState := bucketState); bucketState := bucket.BucketState;
home.M1Status.HomedAndReliable := encoderM1.HomedAndReliable; home.M2Status.HomedAndReliable := encoderM2.HomedAndReliable; home(BucketOffsetValid := bucketState.BucketReferenced, BtnValidation := bench.Operator.JoyBtnRaw);
ADVANCE_TIME(10000000);
bench(M1_PresetTriggerCmd := encoderM1.HwOut.PresetTriggerCmd, M1_PresetValueOut := encoderM1.HwOut.PresetValueOut, M2_PresetTriggerCmd := encoderM2.HwOut.PresetTriggerCmd, M2_PresetValueOut := encoderM2.HwOut.PresetValueOut, RawPosM1 := raw1, RawPosM2 := raw2); raw1 := bench.RawPosM1; raw2 := bench.RawPosM2;
hw1.RawPosIn := bench.Winch.COD1_PosValue; hw1.SlaveOperational := TRUE; hw2.RawPosIn := bench.Winch.COD2_PosValue; hw2.SlaveOperational := TRUE;
encoderM1(Enable := TRUE, HomingPermit := TRUE, HomingAtTargetM := btnM1, CfgHomingTargetM := 8.7, CfgTopSensorPosM := 8.7, HwIn := hw1, Cfg := cfgEncoder, Calib := calibM1); calibM1 := encoderM1.Calib;
bucketEdge(CLK := btnBucket);
encoderM2(Enable := TRUE, HomingPermit := TRUE, HomingAtTargetM := btnM2 OR bucketEdge.Q, CfgHomingTargetM := 23.7, CfgTopSensorPosM := 23.7, UseDynamicTarget := bucketEdge.Q, DynamicHomingTargetM := encoderM1.Measurement.CablePosM + cfgBucket.OffsetCloseM, HwIn := hw2, Cfg := cfgEncoder, Calib := calibM2); calibM2 := encoderM2.Calib;
bucket(Enable := TRUE, Mode := E_Mode.MAINT_N2, PowerContactorEngaged := TRUE, CablePosM1 := encoderM1.Measurement.CablePosM, CablePosM2 := encoderM2.Measurement.CablePosM, HomedM1 := encoderM1.Homed, HomedM2 := encoderM2.Homed, HomedAndReliableM1 := encoderM1.HomedAndReliable, HomedAndReliableM2 := encoderM2.HomedAndReliable, HomingSuspectM1 := encoderM1.HomingSuspect, HomingSuspectM2 := encoderM2.HomingSuspect, ConfirmClosePosition := btnBucket, Config := cfgBucket, BucketState := bucketState); bucketState := bucket.BucketState;
home.M1Status.HomedAndReliable := encoderM1.HomedAndReliable; home.M2Status.HomedAndReliable := encoderM2.HomedAndReliable; home(BucketOffsetValid := bucketState.BucketReferenced, BtnValidation := bench.Operator.JoyBtnRaw);
ASSERT_TRUE(encoderM1.Homed, 'M1 homing accepte'); ASSERT_FALSE(encoderM1.HomingSuspect, 'M1 sans suspicion'); ASSERT_EQ(encoderM1.Fault.ErrorId, 0, 'M1 causes defaut'); ASSERT_FALSE(encoderM1.EncoderFault, 'M1 fiable'); ASSERT_TRUE(encoderM1.HomedAndReliable, 'Premier bouton reference M1'); ASSERT_FALSE(encoderM2.Homed, 'M2 non reference sans son bouton');
btnM2 := TRUE;
ADVANCE_TIME(10000000);
bench(M1_PresetTriggerCmd := encoderM1.HwOut.PresetTriggerCmd, M1_PresetValueOut := encoderM1.HwOut.PresetValueOut, M2_PresetTriggerCmd := encoderM2.HwOut.PresetTriggerCmd, M2_PresetValueOut := encoderM2.HwOut.PresetValueOut, RawPosM1 := raw1, RawPosM2 := raw2); raw1 := bench.RawPosM1; raw2 := bench.RawPosM2;
hw1.RawPosIn := bench.Winch.COD1_PosValue; hw1.SlaveOperational := TRUE; hw2.RawPosIn := bench.Winch.COD2_PosValue; hw2.SlaveOperational := TRUE;
encoderM1(Enable := TRUE, HomingPermit := TRUE, HomingAtTargetM := btnM1, CfgHomingTargetM := 8.7, CfgTopSensorPosM := 8.7, HwIn := hw1, Cfg := cfgEncoder, Calib := calibM1); calibM1 := encoderM1.Calib;
bucketEdge(CLK := btnBucket);
encoderM2(Enable := TRUE, HomingPermit := TRUE, HomingAtTargetM := btnM2 OR bucketEdge.Q, CfgHomingTargetM := 23.7, CfgTopSensorPosM := 23.7, UseDynamicTarget := bucketEdge.Q, DynamicHomingTargetM := encoderM1.Measurement.CablePosM + cfgBucket.OffsetCloseM, HwIn := hw2, Cfg := cfgEncoder, Calib := calibM2); calibM2 := encoderM2.Calib;
bucket(Enable := TRUE, Mode := E_Mode.MAINT_N2, PowerContactorEngaged := TRUE, CablePosM1 := encoderM1.Measurement.CablePosM, CablePosM2 := encoderM2.Measurement.CablePosM, HomedM1 := encoderM1.Homed, HomedM2 := encoderM2.Homed, HomedAndReliableM1 := encoderM1.HomedAndReliable, HomedAndReliableM2 := encoderM2.HomedAndReliable, HomingSuspectM1 := encoderM1.HomingSuspect, HomingSuspectM2 := encoderM2.HomingSuspect, ConfirmClosePosition := btnBucket, Config := cfgBucket, BucketState := bucketState); bucketState := bucket.BucketState;
home.M1Status.HomedAndReliable := encoderM1.HomedAndReliable; home.M2Status.HomedAndReliable := encoderM2.HomedAndReliable; home(BucketOffsetValid := bucketState.BucketReferenced, BtnValidation := bench.Operator.JoyBtnRaw);
btnM2 := FALSE;
ADVANCE_TIME(10000000);
bench(M1_PresetTriggerCmd := encoderM1.HwOut.PresetTriggerCmd, M1_PresetValueOut := encoderM1.HwOut.PresetValueOut, M2_PresetTriggerCmd := encoderM2.HwOut.PresetTriggerCmd, M2_PresetValueOut := encoderM2.HwOut.PresetValueOut, RawPosM1 := raw1, RawPosM2 := raw2); raw1 := bench.RawPosM1; raw2 := bench.RawPosM2;
hw1.RawPosIn := bench.Winch.COD1_PosValue; hw1.SlaveOperational := TRUE; hw2.RawPosIn := bench.Winch.COD2_PosValue; hw2.SlaveOperational := TRUE;
encoderM1(Enable := TRUE, HomingPermit := TRUE, HomingAtTargetM := btnM1, CfgHomingTargetM := 8.7, CfgTopSensorPosM := 8.7, HwIn := hw1, Cfg := cfgEncoder, Calib := calibM1); calibM1 := encoderM1.Calib;
bucketEdge(CLK := btnBucket);
encoderM2(Enable := TRUE, HomingPermit := TRUE, HomingAtTargetM := btnM2 OR bucketEdge.Q, CfgHomingTargetM := 23.7, CfgTopSensorPosM := 23.7, UseDynamicTarget := bucketEdge.Q, DynamicHomingTargetM := encoderM1.Measurement.CablePosM + cfgBucket.OffsetCloseM, HwIn := hw2, Cfg := cfgEncoder, Calib := calibM2); calibM2 := encoderM2.Calib;
bucket(Enable := TRUE, Mode := E_Mode.MAINT_N2, PowerContactorEngaged := TRUE, CablePosM1 := encoderM1.Measurement.CablePosM, CablePosM2 := encoderM2.Measurement.CablePosM, HomedM1 := encoderM1.Homed, HomedM2 := encoderM2.Homed, HomedAndReliableM1 := encoderM1.HomedAndReliable, HomedAndReliableM2 := encoderM2.HomedAndReliable, HomingSuspectM1 := encoderM1.HomingSuspect, HomingSuspectM2 := encoderM2.HomingSuspect, ConfirmClosePosition := btnBucket, Config := cfgBucket, BucketState := bucketState); bucketState := bucket.BucketState;
home.M1Status.HomedAndReliable := encoderM1.HomedAndReliable; home.M2Status.HomedAndReliable := encoderM2.HomedAndReliable; home(BucketOffsetValid := bucketState.BucketReferenced, BtnValidation := bench.Operator.JoyBtnRaw);
ADVANCE_TIME(10000000);
bench(M1_PresetTriggerCmd := encoderM1.HwOut.PresetTriggerCmd, M1_PresetValueOut := encoderM1.HwOut.PresetValueOut, M2_PresetTriggerCmd := encoderM2.HwOut.PresetTriggerCmd, M2_PresetValueOut := encoderM2.HwOut.PresetValueOut, RawPosM1 := raw1, RawPosM2 := raw2); raw1 := bench.RawPosM1; raw2 := bench.RawPosM2;
hw1.RawPosIn := bench.Winch.COD1_PosValue; hw1.SlaveOperational := TRUE; hw2.RawPosIn := bench.Winch.COD2_PosValue; hw2.SlaveOperational := TRUE;
encoderM1(Enable := TRUE, HomingPermit := TRUE, HomingAtTargetM := btnM1, CfgHomingTargetM := 8.7, CfgTopSensorPosM := 8.7, HwIn := hw1, Cfg := cfgEncoder, Calib := calibM1); calibM1 := encoderM1.Calib;
bucketEdge(CLK := btnBucket);
encoderM2(Enable := TRUE, HomingPermit := TRUE, HomingAtTargetM := btnM2 OR bucketEdge.Q, CfgHomingTargetM := 23.7, CfgTopSensorPosM := 23.7, UseDynamicTarget := bucketEdge.Q, DynamicHomingTargetM := encoderM1.Measurement.CablePosM + cfgBucket.OffsetCloseM, HwIn := hw2, Cfg := cfgEncoder, Calib := calibM2); calibM2 := encoderM2.Calib;
bucket(Enable := TRUE, Mode := E_Mode.MAINT_N2, PowerContactorEngaged := TRUE, CablePosM1 := encoderM1.Measurement.CablePosM, CablePosM2 := encoderM2.Measurement.CablePosM, HomedM1 := encoderM1.Homed, HomedM2 := encoderM2.Homed, HomedAndReliableM1 := encoderM1.HomedAndReliable, HomedAndReliableM2 := encoderM2.HomedAndReliable, HomingSuspectM1 := encoderM1.HomingSuspect, HomingSuspectM2 := encoderM2.HomingSuspect, ConfirmClosePosition := btnBucket, Config := cfgBucket, BucketState := bucketState); bucketState := bucket.BucketState;
home.M1Status.HomedAndReliable := encoderM1.HomedAndReliable; home.M2Status.HomedAndReliable := encoderM2.HomedAndReliable; home(BucketOffsetValid := bucketState.BucketReferenced, BtnValidation := bench.Operator.JoyBtnRaw);
ADVANCE_TIME(10000000);
bench(M1_PresetTriggerCmd := encoderM1.HwOut.PresetTriggerCmd, M1_PresetValueOut := encoderM1.HwOut.PresetValueOut, M2_PresetTriggerCmd := encoderM2.HwOut.PresetTriggerCmd, M2_PresetValueOut := encoderM2.HwOut.PresetValueOut, RawPosM1 := raw1, RawPosM2 := raw2); raw1 := bench.RawPosM1; raw2 := bench.RawPosM2;
hw1.RawPosIn := bench.Winch.COD1_PosValue; hw1.SlaveOperational := TRUE; hw2.RawPosIn := bench.Winch.COD2_PosValue; hw2.SlaveOperational := TRUE;
encoderM1(Enable := TRUE, HomingPermit := TRUE, HomingAtTargetM := btnM1, CfgHomingTargetM := 8.7, CfgTopSensorPosM := 8.7, HwIn := hw1, Cfg := cfgEncoder, Calib := calibM1); calibM1 := encoderM1.Calib;
bucketEdge(CLK := btnBucket);
encoderM2(Enable := TRUE, HomingPermit := TRUE, HomingAtTargetM := btnM2 OR bucketEdge.Q, CfgHomingTargetM := 23.7, CfgTopSensorPosM := 23.7, UseDynamicTarget := bucketEdge.Q, DynamicHomingTargetM := encoderM1.Measurement.CablePosM + cfgBucket.OffsetCloseM, HwIn := hw2, Cfg := cfgEncoder, Calib := calibM2); calibM2 := encoderM2.Calib;
bucket(Enable := TRUE, Mode := E_Mode.MAINT_N2, PowerContactorEngaged := TRUE, CablePosM1 := encoderM1.Measurement.CablePosM, CablePosM2 := encoderM2.Measurement.CablePosM, HomedM1 := encoderM1.Homed, HomedM2 := encoderM2.Homed, HomedAndReliableM1 := encoderM1.HomedAndReliable, HomedAndReliableM2 := encoderM2.HomedAndReliable, HomingSuspectM1 := encoderM1.HomingSuspect, HomingSuspectM2 := encoderM2.HomingSuspect, ConfirmClosePosition := btnBucket, Config := cfgBucket, BucketState := bucketState); bucketState := bucket.BucketState;
home.M1Status.HomedAndReliable := encoderM1.HomedAndReliable; home.M2Status.HomedAndReliable := encoderM2.HomedAndReliable; home(BucketOffsetValid := bucketState.BucketReferenced, BtnValidation := bench.Operator.JoyBtnRaw);
ADVANCE_TIME(10000000);
bench(M1_PresetTriggerCmd := encoderM1.HwOut.PresetTriggerCmd, M1_PresetValueOut := encoderM1.HwOut.PresetValueOut, M2_PresetTriggerCmd := encoderM2.HwOut.PresetTriggerCmd, M2_PresetValueOut := encoderM2.HwOut.PresetValueOut, RawPosM1 := raw1, RawPosM2 := raw2); raw1 := bench.RawPosM1; raw2 := bench.RawPosM2;
hw1.RawPosIn := bench.Winch.COD1_PosValue; hw1.SlaveOperational := TRUE; hw2.RawPosIn := bench.Winch.COD2_PosValue; hw2.SlaveOperational := TRUE;
encoderM1(Enable := TRUE, HomingPermit := TRUE, HomingAtTargetM := btnM1, CfgHomingTargetM := 8.7, CfgTopSensorPosM := 8.7, HwIn := hw1, Cfg := cfgEncoder, Calib := calibM1); calibM1 := encoderM1.Calib;
bucketEdge(CLK := btnBucket);
encoderM2(Enable := TRUE, HomingPermit := TRUE, HomingAtTargetM := btnM2 OR bucketEdge.Q, CfgHomingTargetM := 23.7, CfgTopSensorPosM := 23.7, UseDynamicTarget := bucketEdge.Q, DynamicHomingTargetM := encoderM1.Measurement.CablePosM + cfgBucket.OffsetCloseM, HwIn := hw2, Cfg := cfgEncoder, Calib := calibM2); calibM2 := encoderM2.Calib;
bucket(Enable := TRUE, Mode := E_Mode.MAINT_N2, PowerContactorEngaged := TRUE, CablePosM1 := encoderM1.Measurement.CablePosM, CablePosM2 := encoderM2.Measurement.CablePosM, HomedM1 := encoderM1.Homed, HomedM2 := encoderM2.Homed, HomedAndReliableM1 := encoderM1.HomedAndReliable, HomedAndReliableM2 := encoderM2.HomedAndReliable, HomingSuspectM1 := encoderM1.HomingSuspect, HomingSuspectM2 := encoderM2.HomingSuspect, ConfirmClosePosition := btnBucket, Config := cfgBucket, BucketState := bucketState); bucketState := bucket.BucketState;
home.M1Status.HomedAndReliable := encoderM1.HomedAndReliable; home.M2Status.HomedAndReliable := encoderM2.HomedAndReliable; home(BucketOffsetValid := bucketState.BucketReferenced, BtnValidation := bench.Operator.JoyBtnRaw);
ADVANCE_TIME(10000000);
bench(M1_PresetTriggerCmd := encoderM1.HwOut.PresetTriggerCmd, M1_PresetValueOut := encoderM1.HwOut.PresetValueOut, M2_PresetTriggerCmd := encoderM2.HwOut.PresetTriggerCmd, M2_PresetValueOut := encoderM2.HwOut.PresetValueOut, RawPosM1 := raw1, RawPosM2 := raw2); raw1 := bench.RawPosM1; raw2 := bench.RawPosM2;
hw1.RawPosIn := bench.Winch.COD1_PosValue; hw1.SlaveOperational := TRUE; hw2.RawPosIn := bench.Winch.COD2_PosValue; hw2.SlaveOperational := TRUE;
encoderM1(Enable := TRUE, HomingPermit := TRUE, HomingAtTargetM := btnM1, CfgHomingTargetM := 8.7, CfgTopSensorPosM := 8.7, HwIn := hw1, Cfg := cfgEncoder, Calib := calibM1); calibM1 := encoderM1.Calib;
bucketEdge(CLK := btnBucket);
encoderM2(Enable := TRUE, HomingPermit := TRUE, HomingAtTargetM := btnM2 OR bucketEdge.Q, CfgHomingTargetM := 23.7, CfgTopSensorPosM := 23.7, UseDynamicTarget := bucketEdge.Q, DynamicHomingTargetM := encoderM1.Measurement.CablePosM + cfgBucket.OffsetCloseM, HwIn := hw2, Cfg := cfgEncoder, Calib := calibM2); calibM2 := encoderM2.Calib;
bucket(Enable := TRUE, Mode := E_Mode.MAINT_N2, PowerContactorEngaged := TRUE, CablePosM1 := encoderM1.Measurement.CablePosM, CablePosM2 := encoderM2.Measurement.CablePosM, HomedM1 := encoderM1.Homed, HomedM2 := encoderM2.Homed, HomedAndReliableM1 := encoderM1.HomedAndReliable, HomedAndReliableM2 := encoderM2.HomedAndReliable, HomingSuspectM1 := encoderM1.HomingSuspect, HomingSuspectM2 := encoderM2.HomingSuspect, ConfirmClosePosition := btnBucket, Config := cfgBucket, BucketState := bucketState); bucketState := bucket.BucketState;
home.M1Status.HomedAndReliable := encoderM1.HomedAndReliable; home.M2Status.HomedAndReliable := encoderM2.HomedAndReliable; home(BucketOffsetValid := bucketState.BucketReferenced, BtnValidation := bench.Operator.JoyBtnRaw);
ADVANCE_TIME(10000000);
bench(M1_PresetTriggerCmd := encoderM1.HwOut.PresetTriggerCmd, M1_PresetValueOut := encoderM1.HwOut.PresetValueOut, M2_PresetTriggerCmd := encoderM2.HwOut.PresetTriggerCmd, M2_PresetValueOut := encoderM2.HwOut.PresetValueOut, RawPosM1 := raw1, RawPosM2 := raw2); raw1 := bench.RawPosM1; raw2 := bench.RawPosM2;
hw1.RawPosIn := bench.Winch.COD1_PosValue; hw1.SlaveOperational := TRUE; hw2.RawPosIn := bench.Winch.COD2_PosValue; hw2.SlaveOperational := TRUE;
encoderM1(Enable := TRUE, HomingPermit := TRUE, HomingAtTargetM := btnM1, CfgHomingTargetM := 8.7, CfgTopSensorPosM := 8.7, HwIn := hw1, Cfg := cfgEncoder, Calib := calibM1); calibM1 := encoderM1.Calib;
bucketEdge(CLK := btnBucket);
encoderM2(Enable := TRUE, HomingPermit := TRUE, HomingAtTargetM := btnM2 OR bucketEdge.Q, CfgHomingTargetM := 23.7, CfgTopSensorPosM := 23.7, UseDynamicTarget := bucketEdge.Q, DynamicHomingTargetM := encoderM1.Measurement.CablePosM + cfgBucket.OffsetCloseM, HwIn := hw2, Cfg := cfgEncoder, Calib := calibM2); calibM2 := encoderM2.Calib;
bucket(Enable := TRUE, Mode := E_Mode.MAINT_N2, PowerContactorEngaged := TRUE, CablePosM1 := encoderM1.Measurement.CablePosM, CablePosM2 := encoderM2.Measurement.CablePosM, HomedM1 := encoderM1.Homed, HomedM2 := encoderM2.Homed, HomedAndReliableM1 := encoderM1.HomedAndReliable, HomedAndReliableM2 := encoderM2.HomedAndReliable, HomingSuspectM1 := encoderM1.HomingSuspect, HomingSuspectM2 := encoderM2.HomingSuspect, ConfirmClosePosition := btnBucket, Config := cfgBucket, BucketState := bucketState); bucketState := bucket.BucketState;
home.M1Status.HomedAndReliable := encoderM1.HomedAndReliable; home.M2Status.HomedAndReliable := encoderM2.HomedAndReliable; home(BucketOffsetValid := bucketState.BucketReferenced, BtnValidation := bench.Operator.JoyBtnRaw);
ADVANCE_TIME(10000000);
bench(M1_PresetTriggerCmd := encoderM1.HwOut.PresetTriggerCmd, M1_PresetValueOut := encoderM1.HwOut.PresetValueOut, M2_PresetTriggerCmd := encoderM2.HwOut.PresetTriggerCmd, M2_PresetValueOut := encoderM2.HwOut.PresetValueOut, RawPosM1 := raw1, RawPosM2 := raw2); raw1 := bench.RawPosM1; raw2 := bench.RawPosM2;
hw1.RawPosIn := bench.Winch.COD1_PosValue; hw1.SlaveOperational := TRUE; hw2.RawPosIn := bench.Winch.COD2_PosValue; hw2.SlaveOperational := TRUE;
encoderM1(Enable := TRUE, HomingPermit := TRUE, HomingAtTargetM := btnM1, CfgHomingTargetM := 8.7, CfgTopSensorPosM := 8.7, HwIn := hw1, Cfg := cfgEncoder, Calib := calibM1); calibM1 := encoderM1.Calib;
bucketEdge(CLK := btnBucket);
encoderM2(Enable := TRUE, HomingPermit := TRUE, HomingAtTargetM := btnM2 OR bucketEdge.Q, CfgHomingTargetM := 23.7, CfgTopSensorPosM := 23.7, UseDynamicTarget := bucketEdge.Q, DynamicHomingTargetM := encoderM1.Measurement.CablePosM + cfgBucket.OffsetCloseM, HwIn := hw2, Cfg := cfgEncoder, Calib := calibM2); calibM2 := encoderM2.Calib;
bucket(Enable := TRUE, Mode := E_Mode.MAINT_N2, PowerContactorEngaged := TRUE, CablePosM1 := encoderM1.Measurement.CablePosM, CablePosM2 := encoderM2.Measurement.CablePosM, HomedM1 := encoderM1.Homed, HomedM2 := encoderM2.Homed, HomedAndReliableM1 := encoderM1.HomedAndReliable, HomedAndReliableM2 := encoderM2.HomedAndReliable, HomingSuspectM1 := encoderM1.HomingSuspect, HomingSuspectM2 := encoderM2.HomingSuspect, ConfirmClosePosition := btnBucket, Config := cfgBucket, BucketState := bucketState); bucketState := bucket.BucketState;
home.M1Status.HomedAndReliable := encoderM1.HomedAndReliable; home.M2Status.HomedAndReliable := encoderM2.HomedAndReliable; home(BucketOffsetValid := bucketState.BucketReferenced, BtnValidation := bench.Operator.JoyBtnRaw);
ADVANCE_TIME(10000000);
bench(M1_PresetTriggerCmd := encoderM1.HwOut.PresetTriggerCmd, M1_PresetValueOut := encoderM1.HwOut.PresetValueOut, M2_PresetTriggerCmd := encoderM2.HwOut.PresetTriggerCmd, M2_PresetValueOut := encoderM2.HwOut.PresetValueOut, RawPosM1 := raw1, RawPosM2 := raw2); raw1 := bench.RawPosM1; raw2 := bench.RawPosM2;
hw1.RawPosIn := bench.Winch.COD1_PosValue; hw1.SlaveOperational := TRUE; hw2.RawPosIn := bench.Winch.COD2_PosValue; hw2.SlaveOperational := TRUE;
encoderM1(Enable := TRUE, HomingPermit := TRUE, HomingAtTargetM := btnM1, CfgHomingTargetM := 8.7, CfgTopSensorPosM := 8.7, HwIn := hw1, Cfg := cfgEncoder, Calib := calibM1); calibM1 := encoderM1.Calib;
bucketEdge(CLK := btnBucket);
encoderM2(Enable := TRUE, HomingPermit := TRUE, HomingAtTargetM := btnM2 OR bucketEdge.Q, CfgHomingTargetM := 23.7, CfgTopSensorPosM := 23.7, UseDynamicTarget := bucketEdge.Q, DynamicHomingTargetM := encoderM1.Measurement.CablePosM + cfgBucket.OffsetCloseM, HwIn := hw2, Cfg := cfgEncoder, Calib := calibM2); calibM2 := encoderM2.Calib;
bucket(Enable := TRUE, Mode := E_Mode.MAINT_N2, PowerContactorEngaged := TRUE, CablePosM1 := encoderM1.Measurement.CablePosM, CablePosM2 := encoderM2.Measurement.CablePosM, HomedM1 := encoderM1.Homed, HomedM2 := encoderM2.Homed, HomedAndReliableM1 := encoderM1.HomedAndReliable, HomedAndReliableM2 := encoderM2.HomedAndReliable, HomingSuspectM1 := encoderM1.HomingSuspect, HomingSuspectM2 := encoderM2.HomingSuspect, ConfirmClosePosition := btnBucket, Config := cfgBucket, BucketState := bucketState); bucketState := bucket.BucketState;
home.M1Status.HomedAndReliable := encoderM1.HomedAndReliable; home.M2Status.HomedAndReliable := encoderM2.HomedAndReliable; home(BucketOffsetValid := bucketState.BucketReferenced, BtnValidation := bench.Operator.JoyBtnRaw);
ADVANCE_TIME(10000000);
bench(M1_PresetTriggerCmd := encoderM1.HwOut.PresetTriggerCmd, M1_PresetValueOut := encoderM1.HwOut.PresetValueOut, M2_PresetTriggerCmd := encoderM2.HwOut.PresetTriggerCmd, M2_PresetValueOut := encoderM2.HwOut.PresetValueOut, RawPosM1 := raw1, RawPosM2 := raw2); raw1 := bench.RawPosM1; raw2 := bench.RawPosM2;
hw1.RawPosIn := bench.Winch.COD1_PosValue; hw1.SlaveOperational := TRUE; hw2.RawPosIn := bench.Winch.COD2_PosValue; hw2.SlaveOperational := TRUE;
encoderM1(Enable := TRUE, HomingPermit := TRUE, HomingAtTargetM := btnM1, CfgHomingTargetM := 8.7, CfgTopSensorPosM := 8.7, HwIn := hw1, Cfg := cfgEncoder, Calib := calibM1); calibM1 := encoderM1.Calib;
bucketEdge(CLK := btnBucket);
encoderM2(Enable := TRUE, HomingPermit := TRUE, HomingAtTargetM := btnM2 OR bucketEdge.Q, CfgHomingTargetM := 23.7, CfgTopSensorPosM := 23.7, UseDynamicTarget := bucketEdge.Q, DynamicHomingTargetM := encoderM1.Measurement.CablePosM + cfgBucket.OffsetCloseM, HwIn := hw2, Cfg := cfgEncoder, Calib := calibM2); calibM2 := encoderM2.Calib;
bucket(Enable := TRUE, Mode := E_Mode.MAINT_N2, PowerContactorEngaged := TRUE, CablePosM1 := encoderM1.Measurement.CablePosM, CablePosM2 := encoderM2.Measurement.CablePosM, HomedM1 := encoderM1.Homed, HomedM2 := encoderM2.Homed, HomedAndReliableM1 := encoderM1.HomedAndReliable, HomedAndReliableM2 := encoderM2.HomedAndReliable, HomingSuspectM1 := encoderM1.HomingSuspect, HomingSuspectM2 := encoderM2.HomingSuspect, ConfirmClosePosition := btnBucket, Config := cfgBucket, BucketState := bucketState); bucketState := bucket.BucketState;
home.M1Status.HomedAndReliable := encoderM1.HomedAndReliable; home.M2Status.HomedAndReliable := encoderM2.HomedAndReliable; home(BucketOffsetValid := bucketState.BucketReferenced, BtnValidation := bench.Operator.JoyBtnRaw);
ADVANCE_TIME(10000000);
bench(M1_PresetTriggerCmd := encoderM1.HwOut.PresetTriggerCmd, M1_PresetValueOut := encoderM1.HwOut.PresetValueOut, M2_PresetTriggerCmd := encoderM2.HwOut.PresetTriggerCmd, M2_PresetValueOut := encoderM2.HwOut.PresetValueOut, RawPosM1 := raw1, RawPosM2 := raw2); raw1 := bench.RawPosM1; raw2 := bench.RawPosM2;
hw1.RawPosIn := bench.Winch.COD1_PosValue; hw1.SlaveOperational := TRUE; hw2.RawPosIn := bench.Winch.COD2_PosValue; hw2.SlaveOperational := TRUE;
encoderM1(Enable := TRUE, HomingPermit := TRUE, HomingAtTargetM := btnM1, CfgHomingTargetM := 8.7, CfgTopSensorPosM := 8.7, HwIn := hw1, Cfg := cfgEncoder, Calib := calibM1); calibM1 := encoderM1.Calib;
bucketEdge(CLK := btnBucket);
encoderM2(Enable := TRUE, HomingPermit := TRUE, HomingAtTargetM := btnM2 OR bucketEdge.Q, CfgHomingTargetM := 23.7, CfgTopSensorPosM := 23.7, UseDynamicTarget := bucketEdge.Q, DynamicHomingTargetM := encoderM1.Measurement.CablePosM + cfgBucket.OffsetCloseM, HwIn := hw2, Cfg := cfgEncoder, Calib := calibM2); calibM2 := encoderM2.Calib;
bucket(Enable := TRUE, Mode := E_Mode.MAINT_N2, PowerContactorEngaged := TRUE, CablePosM1 := encoderM1.Measurement.CablePosM, CablePosM2 := encoderM2.Measurement.CablePosM, HomedM1 := encoderM1.Homed, HomedM2 := encoderM2.Homed, HomedAndReliableM1 := encoderM1.HomedAndReliable, HomedAndReliableM2 := encoderM2.HomedAndReliable, HomingSuspectM1 := encoderM1.HomingSuspect, HomingSuspectM2 := encoderM2.HomingSuspect, ConfirmClosePosition := btnBucket, Config := cfgBucket, BucketState := bucketState); bucketState := bucket.BucketState;
home.M1Status.HomedAndReliable := encoderM1.HomedAndReliable; home.M2Status.HomedAndReliable := encoderM2.HomedAndReliable; home(BucketOffsetValid := bucketState.BucketReferenced, BtnValidation := bench.Operator.JoyBtnRaw);
ADVANCE_TIME(10000000);
bench(M1_PresetTriggerCmd := encoderM1.HwOut.PresetTriggerCmd, M1_PresetValueOut := encoderM1.HwOut.PresetValueOut, M2_PresetTriggerCmd := encoderM2.HwOut.PresetTriggerCmd, M2_PresetValueOut := encoderM2.HwOut.PresetValueOut, RawPosM1 := raw1, RawPosM2 := raw2); raw1 := bench.RawPosM1; raw2 := bench.RawPosM2;
hw1.RawPosIn := bench.Winch.COD1_PosValue; hw1.SlaveOperational := TRUE; hw2.RawPosIn := bench.Winch.COD2_PosValue; hw2.SlaveOperational := TRUE;
encoderM1(Enable := TRUE, HomingPermit := TRUE, HomingAtTargetM := btnM1, CfgHomingTargetM := 8.7, CfgTopSensorPosM := 8.7, HwIn := hw1, Cfg := cfgEncoder, Calib := calibM1); calibM1 := encoderM1.Calib;
bucketEdge(CLK := btnBucket);
encoderM2(Enable := TRUE, HomingPermit := TRUE, HomingAtTargetM := btnM2 OR bucketEdge.Q, CfgHomingTargetM := 23.7, CfgTopSensorPosM := 23.7, UseDynamicTarget := bucketEdge.Q, DynamicHomingTargetM := encoderM1.Measurement.CablePosM + cfgBucket.OffsetCloseM, HwIn := hw2, Cfg := cfgEncoder, Calib := calibM2); calibM2 := encoderM2.Calib;
bucket(Enable := TRUE, Mode := E_Mode.MAINT_N2, PowerContactorEngaged := TRUE, CablePosM1 := encoderM1.Measurement.CablePosM, CablePosM2 := encoderM2.Measurement.CablePosM, HomedM1 := encoderM1.Homed, HomedM2 := encoderM2.Homed, HomedAndReliableM1 := encoderM1.HomedAndReliable, HomedAndReliableM2 := encoderM2.HomedAndReliable, HomingSuspectM1 := encoderM1.HomingSuspect, HomingSuspectM2 := encoderM2.HomingSuspect, ConfirmClosePosition := btnBucket, Config := cfgBucket, BucketState := bucketState); bucketState := bucket.BucketState;
home.M1Status.HomedAndReliable := encoderM1.HomedAndReliable; home.M2Status.HomedAndReliable := encoderM2.HomedAndReliable; home(BucketOffsetValid := bucketState.BucketReferenced, BtnValidation := bench.Operator.JoyBtnRaw);
ADVANCE_TIME(10000000);
bench(M1_PresetTriggerCmd := encoderM1.HwOut.PresetTriggerCmd, M1_PresetValueOut := encoderM1.HwOut.PresetValueOut, M2_PresetTriggerCmd := encoderM2.HwOut.PresetTriggerCmd, M2_PresetValueOut := encoderM2.HwOut.PresetValueOut, RawPosM1 := raw1, RawPosM2 := raw2); raw1 := bench.RawPosM1; raw2 := bench.RawPosM2;
hw1.RawPosIn := bench.Winch.COD1_PosValue; hw1.SlaveOperational := TRUE; hw2.RawPosIn := bench.Winch.COD2_PosValue; hw2.SlaveOperational := TRUE;
encoderM1(Enable := TRUE, HomingPermit := TRUE, HomingAtTargetM := btnM1, CfgHomingTargetM := 8.7, CfgTopSensorPosM := 8.7, HwIn := hw1, Cfg := cfgEncoder, Calib := calibM1); calibM1 := encoderM1.Calib;
bucketEdge(CLK := btnBucket);
encoderM2(Enable := TRUE, HomingPermit := TRUE, HomingAtTargetM := btnM2 OR bucketEdge.Q, CfgHomingTargetM := 23.7, CfgTopSensorPosM := 23.7, UseDynamicTarget := bucketEdge.Q, DynamicHomingTargetM := encoderM1.Measurement.CablePosM + cfgBucket.OffsetCloseM, HwIn := hw2, Cfg := cfgEncoder, Calib := calibM2); calibM2 := encoderM2.Calib;
bucket(Enable := TRUE, Mode := E_Mode.MAINT_N2, PowerContactorEngaged := TRUE, CablePosM1 := encoderM1.Measurement.CablePosM, CablePosM2 := encoderM2.Measurement.CablePosM, HomedM1 := encoderM1.Homed, HomedM2 := encoderM2.Homed, HomedAndReliableM1 := encoderM1.HomedAndReliable, HomedAndReliableM2 := encoderM2.HomedAndReliable, HomingSuspectM1 := encoderM1.HomingSuspect, HomingSuspectM2 := encoderM2.HomingSuspect, ConfirmClosePosition := btnBucket, Config := cfgBucket, BucketState := bucketState); bucketState := bucket.BucketState;
home.M1Status.HomedAndReliable := encoderM1.HomedAndReliable; home.M2Status.HomedAndReliable := encoderM2.HomedAndReliable; home(BucketOffsetValid := bucketState.BucketReferenced, BtnValidation := bench.Operator.JoyBtnRaw);
ADVANCE_TIME(10000000);
bench(M1_PresetTriggerCmd := encoderM1.HwOut.PresetTriggerCmd, M1_PresetValueOut := encoderM1.HwOut.PresetValueOut, M2_PresetTriggerCmd := encoderM2.HwOut.PresetTriggerCmd, M2_PresetValueOut := encoderM2.HwOut.PresetValueOut, RawPosM1 := raw1, RawPosM2 := raw2); raw1 := bench.RawPosM1; raw2 := bench.RawPosM2;
hw1.RawPosIn := bench.Winch.COD1_PosValue; hw1.SlaveOperational := TRUE; hw2.RawPosIn := bench.Winch.COD2_PosValue; hw2.SlaveOperational := TRUE;
encoderM1(Enable := TRUE, HomingPermit := TRUE, HomingAtTargetM := btnM1, CfgHomingTargetM := 8.7, CfgTopSensorPosM := 8.7, HwIn := hw1, Cfg := cfgEncoder, Calib := calibM1); calibM1 := encoderM1.Calib;
bucketEdge(CLK := btnBucket);
encoderM2(Enable := TRUE, HomingPermit := TRUE, HomingAtTargetM := btnM2 OR bucketEdge.Q, CfgHomingTargetM := 23.7, CfgTopSensorPosM := 23.7, UseDynamicTarget := bucketEdge.Q, DynamicHomingTargetM := encoderM1.Measurement.CablePosM + cfgBucket.OffsetCloseM, HwIn := hw2, Cfg := cfgEncoder, Calib := calibM2); calibM2 := encoderM2.Calib;
bucket(Enable := TRUE, Mode := E_Mode.MAINT_N2, PowerContactorEngaged := TRUE, CablePosM1 := encoderM1.Measurement.CablePosM, CablePosM2 := encoderM2.Measurement.CablePosM, HomedM1 := encoderM1.Homed, HomedM2 := encoderM2.Homed, HomedAndReliableM1 := encoderM1.HomedAndReliable, HomedAndReliableM2 := encoderM2.HomedAndReliable, HomingSuspectM1 := encoderM1.HomingSuspect, HomingSuspectM2 := encoderM2.HomingSuspect, ConfirmClosePosition := btnBucket, Config := cfgBucket, BucketState := bucketState); bucketState := bucket.BucketState;
home.M1Status.HomedAndReliable := encoderM1.HomedAndReliable; home.M2Status.HomedAndReliable := encoderM2.HomedAndReliable; home(BucketOffsetValid := bucketState.BucketReferenced, BtnValidation := bench.Operator.JoyBtnRaw);
ADVANCE_TIME(10000000);
bench(M1_PresetTriggerCmd := encoderM1.HwOut.PresetTriggerCmd, M1_PresetValueOut := encoderM1.HwOut.PresetValueOut, M2_PresetTriggerCmd := encoderM2.HwOut.PresetTriggerCmd, M2_PresetValueOut := encoderM2.HwOut.PresetValueOut, RawPosM1 := raw1, RawPosM2 := raw2); raw1 := bench.RawPosM1; raw2 := bench.RawPosM2;
hw1.RawPosIn := bench.Winch.COD1_PosValue; hw1.SlaveOperational := TRUE; hw2.RawPosIn := bench.Winch.COD2_PosValue; hw2.SlaveOperational := TRUE;
encoderM1(Enable := TRUE, HomingPermit := TRUE, HomingAtTargetM := btnM1, CfgHomingTargetM := 8.7, CfgTopSensorPosM := 8.7, HwIn := hw1, Cfg := cfgEncoder, Calib := calibM1); calibM1 := encoderM1.Calib;
bucketEdge(CLK := btnBucket);
encoderM2(Enable := TRUE, HomingPermit := TRUE, HomingAtTargetM := btnM2 OR bucketEdge.Q, CfgHomingTargetM := 23.7, CfgTopSensorPosM := 23.7, UseDynamicTarget := bucketEdge.Q, DynamicHomingTargetM := encoderM1.Measurement.CablePosM + cfgBucket.OffsetCloseM, HwIn := hw2, Cfg := cfgEncoder, Calib := calibM2); calibM2 := encoderM2.Calib;
bucket(Enable := TRUE, Mode := E_Mode.MAINT_N2, PowerContactorEngaged := TRUE, CablePosM1 := encoderM1.Measurement.CablePosM, CablePosM2 := encoderM2.Measurement.CablePosM, HomedM1 := encoderM1.Homed, HomedM2 := encoderM2.Homed, HomedAndReliableM1 := encoderM1.HomedAndReliable, HomedAndReliableM2 := encoderM2.HomedAndReliable, HomingSuspectM1 := encoderM1.HomingSuspect, HomingSuspectM2 := encoderM2.HomingSuspect, ConfirmClosePosition := btnBucket, Config := cfgBucket, BucketState := bucketState); bucketState := bucket.BucketState;
home.M1Status.HomedAndReliable := encoderM1.HomedAndReliable; home.M2Status.HomedAndReliable := encoderM2.HomedAndReliable; home(BucketOffsetValid := bucketState.BucketReferenced, BtnValidation := bench.Operator.JoyBtnRaw);
ADVANCE_TIME(10000000);
bench(M1_PresetTriggerCmd := encoderM1.HwOut.PresetTriggerCmd, M1_PresetValueOut := encoderM1.HwOut.PresetValueOut, M2_PresetTriggerCmd := encoderM2.HwOut.PresetTriggerCmd, M2_PresetValueOut := encoderM2.HwOut.PresetValueOut, RawPosM1 := raw1, RawPosM2 := raw2); raw1 := bench.RawPosM1; raw2 := bench.RawPosM2;
hw1.RawPosIn := bench.Winch.COD1_PosValue; hw1.SlaveOperational := TRUE; hw2.RawPosIn := bench.Winch.COD2_PosValue; hw2.SlaveOperational := TRUE;
encoderM1(Enable := TRUE, HomingPermit := TRUE, HomingAtTargetM := btnM1, CfgHomingTargetM := 8.7, CfgTopSensorPosM := 8.7, HwIn := hw1, Cfg := cfgEncoder, Calib := calibM1); calibM1 := encoderM1.Calib;
bucketEdge(CLK := btnBucket);
encoderM2(Enable := TRUE, HomingPermit := TRUE, HomingAtTargetM := btnM2 OR bucketEdge.Q, CfgHomingTargetM := 23.7, CfgTopSensorPosM := 23.7, UseDynamicTarget := bucketEdge.Q, DynamicHomingTargetM := encoderM1.Measurement.CablePosM + cfgBucket.OffsetCloseM, HwIn := hw2, Cfg := cfgEncoder, Calib := calibM2); calibM2 := encoderM2.Calib;
bucket(Enable := TRUE, Mode := E_Mode.MAINT_N2, PowerContactorEngaged := TRUE, CablePosM1 := encoderM1.Measurement.CablePosM, CablePosM2 := encoderM2.Measurement.CablePosM, HomedM1 := encoderM1.Homed, HomedM2 := encoderM2.Homed, HomedAndReliableM1 := encoderM1.HomedAndReliable, HomedAndReliableM2 := encoderM2.HomedAndReliable, HomingSuspectM1 := encoderM1.HomingSuspect, HomingSuspectM2 := encoderM2.HomingSuspect, ConfirmClosePosition := btnBucket, Config := cfgBucket, BucketState := bucketState); bucketState := bucket.BucketState;
home.M1Status.HomedAndReliable := encoderM1.HomedAndReliable; home.M2Status.HomedAndReliable := encoderM2.HomedAndReliable; home(BucketOffsetValid := bucketState.BucketReferenced, BtnValidation := bench.Operator.JoyBtnRaw);
ADVANCE_TIME(10000000);
bench(M1_PresetTriggerCmd := encoderM1.HwOut.PresetTriggerCmd, M1_PresetValueOut := encoderM1.HwOut.PresetValueOut, M2_PresetTriggerCmd := encoderM2.HwOut.PresetTriggerCmd, M2_PresetValueOut := encoderM2.HwOut.PresetValueOut, RawPosM1 := raw1, RawPosM2 := raw2); raw1 := bench.RawPosM1; raw2 := bench.RawPosM2;
hw1.RawPosIn := bench.Winch.COD1_PosValue; hw1.SlaveOperational := TRUE; hw2.RawPosIn := bench.Winch.COD2_PosValue; hw2.SlaveOperational := TRUE;
encoderM1(Enable := TRUE, HomingPermit := TRUE, HomingAtTargetM := btnM1, CfgHomingTargetM := 8.7, CfgTopSensorPosM := 8.7, HwIn := hw1, Cfg := cfgEncoder, Calib := calibM1); calibM1 := encoderM1.Calib;
bucketEdge(CLK := btnBucket);
encoderM2(Enable := TRUE, HomingPermit := TRUE, HomingAtTargetM := btnM2 OR bucketEdge.Q, CfgHomingTargetM := 23.7, CfgTopSensorPosM := 23.7, UseDynamicTarget := bucketEdge.Q, DynamicHomingTargetM := encoderM1.Measurement.CablePosM + cfgBucket.OffsetCloseM, HwIn := hw2, Cfg := cfgEncoder, Calib := calibM2); calibM2 := encoderM2.Calib;
bucket(Enable := TRUE, Mode := E_Mode.MAINT_N2, PowerContactorEngaged := TRUE, CablePosM1 := encoderM1.Measurement.CablePosM, CablePosM2 := encoderM2.Measurement.CablePosM, HomedM1 := encoderM1.Homed, HomedM2 := encoderM2.Homed, HomedAndReliableM1 := encoderM1.HomedAndReliable, HomedAndReliableM2 := encoderM2.HomedAndReliable, HomingSuspectM1 := encoderM1.HomingSuspect, HomingSuspectM2 := encoderM2.HomingSuspect, ConfirmClosePosition := btnBucket, Config := cfgBucket, BucketState := bucketState); bucketState := bucket.BucketState;
home.M1Status.HomedAndReliable := encoderM1.HomedAndReliable; home.M2Status.HomedAndReliable := encoderM2.HomedAndReliable; home(BucketOffsetValid := bucketState.BucketReferenced, BtnValidation := bench.Operator.JoyBtnRaw);
ADVANCE_TIME(10000000);
bench(M1_PresetTriggerCmd := encoderM1.HwOut.PresetTriggerCmd, M1_PresetValueOut := encoderM1.HwOut.PresetValueOut, M2_PresetTriggerCmd := encoderM2.HwOut.PresetTriggerCmd, M2_PresetValueOut := encoderM2.HwOut.PresetValueOut, RawPosM1 := raw1, RawPosM2 := raw2); raw1 := bench.RawPosM1; raw2 := bench.RawPosM2;
hw1.RawPosIn := bench.Winch.COD1_PosValue; hw1.SlaveOperational := TRUE; hw2.RawPosIn := bench.Winch.COD2_PosValue; hw2.SlaveOperational := TRUE;
encoderM1(Enable := TRUE, HomingPermit := TRUE, HomingAtTargetM := btnM1, CfgHomingTargetM := 8.7, CfgTopSensorPosM := 8.7, HwIn := hw1, Cfg := cfgEncoder, Calib := calibM1); calibM1 := encoderM1.Calib;
bucketEdge(CLK := btnBucket);
encoderM2(Enable := TRUE, HomingPermit := TRUE, HomingAtTargetM := btnM2 OR bucketEdge.Q, CfgHomingTargetM := 23.7, CfgTopSensorPosM := 23.7, UseDynamicTarget := bucketEdge.Q, DynamicHomingTargetM := encoderM1.Measurement.CablePosM + cfgBucket.OffsetCloseM, HwIn := hw2, Cfg := cfgEncoder, Calib := calibM2); calibM2 := encoderM2.Calib;
bucket(Enable := TRUE, Mode := E_Mode.MAINT_N2, PowerContactorEngaged := TRUE, CablePosM1 := encoderM1.Measurement.CablePosM, CablePosM2 := encoderM2.Measurement.CablePosM, HomedM1 := encoderM1.Homed, HomedM2 := encoderM2.Homed, HomedAndReliableM1 := encoderM1.HomedAndReliable, HomedAndReliableM2 := encoderM2.HomedAndReliable, HomingSuspectM1 := encoderM1.HomingSuspect, HomingSuspectM2 := encoderM2.HomingSuspect, ConfirmClosePosition := btnBucket, Config := cfgBucket, BucketState := bucketState); bucketState := bucket.BucketState;
home.M1Status.HomedAndReliable := encoderM1.HomedAndReliable; home.M2Status.HomedAndReliable := encoderM2.HomedAndReliable; home(BucketOffsetValid := bucketState.BucketReferenced, BtnValidation := bench.Operator.JoyBtnRaw);
ADVANCE_TIME(10000000);
bench(M1_PresetTriggerCmd := encoderM1.HwOut.PresetTriggerCmd, M1_PresetValueOut := encoderM1.HwOut.PresetValueOut, M2_PresetTriggerCmd := encoderM2.HwOut.PresetTriggerCmd, M2_PresetValueOut := encoderM2.HwOut.PresetValueOut, RawPosM1 := raw1, RawPosM2 := raw2); raw1 := bench.RawPosM1; raw2 := bench.RawPosM2;
hw1.RawPosIn := bench.Winch.COD1_PosValue; hw1.SlaveOperational := TRUE; hw2.RawPosIn := bench.Winch.COD2_PosValue; hw2.SlaveOperational := TRUE;
encoderM1(Enable := TRUE, HomingPermit := TRUE, HomingAtTargetM := btnM1, CfgHomingTargetM := 8.7, CfgTopSensorPosM := 8.7, HwIn := hw1, Cfg := cfgEncoder, Calib := calibM1); calibM1 := encoderM1.Calib;
bucketEdge(CLK := btnBucket);
encoderM2(Enable := TRUE, HomingPermit := TRUE, HomingAtTargetM := btnM2 OR bucketEdge.Q, CfgHomingTargetM := 23.7, CfgTopSensorPosM := 23.7, UseDynamicTarget := bucketEdge.Q, DynamicHomingTargetM := encoderM1.Measurement.CablePosM + cfgBucket.OffsetCloseM, HwIn := hw2, Cfg := cfgEncoder, Calib := calibM2); calibM2 := encoderM2.Calib;
bucket(Enable := TRUE, Mode := E_Mode.MAINT_N2, PowerContactorEngaged := TRUE, CablePosM1 := encoderM1.Measurement.CablePosM, CablePosM2 := encoderM2.Measurement.CablePosM, HomedM1 := encoderM1.Homed, HomedM2 := encoderM2.Homed, HomedAndReliableM1 := encoderM1.HomedAndReliable, HomedAndReliableM2 := encoderM2.HomedAndReliable, HomingSuspectM1 := encoderM1.HomingSuspect, HomingSuspectM2 := encoderM2.HomingSuspect, ConfirmClosePosition := btnBucket, Config := cfgBucket, BucketState := bucketState); bucketState := bucket.BucketState;
home.M1Status.HomedAndReliable := encoderM1.HomedAndReliable; home.M2Status.HomedAndReliable := encoderM2.HomedAndReliable; home(BucketOffsetValid := bucketState.BucketReferenced, BtnValidation := bench.Operator.JoyBtnRaw);
ADVANCE_TIME(10000000);
bench(M1_PresetTriggerCmd := encoderM1.HwOut.PresetTriggerCmd, M1_PresetValueOut := encoderM1.HwOut.PresetValueOut, M2_PresetTriggerCmd := encoderM2.HwOut.PresetTriggerCmd, M2_PresetValueOut := encoderM2.HwOut.PresetValueOut, RawPosM1 := raw1, RawPosM2 := raw2); raw1 := bench.RawPosM1; raw2 := bench.RawPosM2;
hw1.RawPosIn := bench.Winch.COD1_PosValue; hw1.SlaveOperational := TRUE; hw2.RawPosIn := bench.Winch.COD2_PosValue; hw2.SlaveOperational := TRUE;
encoderM1(Enable := TRUE, HomingPermit := TRUE, HomingAtTargetM := btnM1, CfgHomingTargetM := 8.7, CfgTopSensorPosM := 8.7, HwIn := hw1, Cfg := cfgEncoder, Calib := calibM1); calibM1 := encoderM1.Calib;
bucketEdge(CLK := btnBucket);
encoderM2(Enable := TRUE, HomingPermit := TRUE, HomingAtTargetM := btnM2 OR bucketEdge.Q, CfgHomingTargetM := 23.7, CfgTopSensorPosM := 23.7, UseDynamicTarget := bucketEdge.Q, DynamicHomingTargetM := encoderM1.Measurement.CablePosM + cfgBucket.OffsetCloseM, HwIn := hw2, Cfg := cfgEncoder, Calib := calibM2); calibM2 := encoderM2.Calib;
bucket(Enable := TRUE, Mode := E_Mode.MAINT_N2, PowerContactorEngaged := TRUE, CablePosM1 := encoderM1.Measurement.CablePosM, CablePosM2 := encoderM2.Measurement.CablePosM, HomedM1 := encoderM1.Homed, HomedM2 := encoderM2.Homed, HomedAndReliableM1 := encoderM1.HomedAndReliable, HomedAndReliableM2 := encoderM2.HomedAndReliable, HomingSuspectM1 := encoderM1.HomingSuspect, HomingSuspectM2 := encoderM2.HomingSuspect, ConfirmClosePosition := btnBucket, Config := cfgBucket, BucketState := bucketState); bucketState := bucket.BucketState;
home.M1Status.HomedAndReliable := encoderM1.HomedAndReliable; home.M2Status.HomedAndReliable := encoderM2.HomedAndReliable; home(BucketOffsetValid := bucketState.BucketReferenced, BtnValidation := bench.Operator.JoyBtnRaw);
ADVANCE_TIME(10000000);
bench(M1_PresetTriggerCmd := encoderM1.HwOut.PresetTriggerCmd, M1_PresetValueOut := encoderM1.HwOut.PresetValueOut, M2_PresetTriggerCmd := encoderM2.HwOut.PresetTriggerCmd, M2_PresetValueOut := encoderM2.HwOut.PresetValueOut, RawPosM1 := raw1, RawPosM2 := raw2); raw1 := bench.RawPosM1; raw2 := bench.RawPosM2;
hw1.RawPosIn := bench.Winch.COD1_PosValue; hw1.SlaveOperational := TRUE; hw2.RawPosIn := bench.Winch.COD2_PosValue; hw2.SlaveOperational := TRUE;
encoderM1(Enable := TRUE, HomingPermit := TRUE, HomingAtTargetM := btnM1, CfgHomingTargetM := 8.7, CfgTopSensorPosM := 8.7, HwIn := hw1, Cfg := cfgEncoder, Calib := calibM1); calibM1 := encoderM1.Calib;
bucketEdge(CLK := btnBucket);
encoderM2(Enable := TRUE, HomingPermit := TRUE, HomingAtTargetM := btnM2 OR bucketEdge.Q, CfgHomingTargetM := 23.7, CfgTopSensorPosM := 23.7, UseDynamicTarget := bucketEdge.Q, DynamicHomingTargetM := encoderM1.Measurement.CablePosM + cfgBucket.OffsetCloseM, HwIn := hw2, Cfg := cfgEncoder, Calib := calibM2); calibM2 := encoderM2.Calib;
bucket(Enable := TRUE, Mode := E_Mode.MAINT_N2, PowerContactorEngaged := TRUE, CablePosM1 := encoderM1.Measurement.CablePosM, CablePosM2 := encoderM2.Measurement.CablePosM, HomedM1 := encoderM1.Homed, HomedM2 := encoderM2.Homed, HomedAndReliableM1 := encoderM1.HomedAndReliable, HomedAndReliableM2 := encoderM2.HomedAndReliable, HomingSuspectM1 := encoderM1.HomingSuspect, HomingSuspectM2 := encoderM2.HomingSuspect, ConfirmClosePosition := btnBucket, Config := cfgBucket, BucketState := bucketState); bucketState := bucket.BucketState;
home.M1Status.HomedAndReliable := encoderM1.HomedAndReliable; home.M2Status.HomedAndReliable := encoderM2.HomedAndReliable; home(BucketOffsetValid := bucketState.BucketReferenced, BtnValidation := bench.Operator.JoyBtnRaw);
ADVANCE_TIME(10000000);
bench(M1_PresetTriggerCmd := encoderM1.HwOut.PresetTriggerCmd, M1_PresetValueOut := encoderM1.HwOut.PresetValueOut, M2_PresetTriggerCmd := encoderM2.HwOut.PresetTriggerCmd, M2_PresetValueOut := encoderM2.HwOut.PresetValueOut, RawPosM1 := raw1, RawPosM2 := raw2); raw1 := bench.RawPosM1; raw2 := bench.RawPosM2;
hw1.RawPosIn := bench.Winch.COD1_PosValue; hw1.SlaveOperational := TRUE; hw2.RawPosIn := bench.Winch.COD2_PosValue; hw2.SlaveOperational := TRUE;
encoderM1(Enable := TRUE, HomingPermit := TRUE, HomingAtTargetM := btnM1, CfgHomingTargetM := 8.7, CfgTopSensorPosM := 8.7, HwIn := hw1, Cfg := cfgEncoder, Calib := calibM1); calibM1 := encoderM1.Calib;
bucketEdge(CLK := btnBucket);
encoderM2(Enable := TRUE, HomingPermit := TRUE, HomingAtTargetM := btnM2 OR bucketEdge.Q, CfgHomingTargetM := 23.7, CfgTopSensorPosM := 23.7, UseDynamicTarget := bucketEdge.Q, DynamicHomingTargetM := encoderM1.Measurement.CablePosM + cfgBucket.OffsetCloseM, HwIn := hw2, Cfg := cfgEncoder, Calib := calibM2); calibM2 := encoderM2.Calib;
bucket(Enable := TRUE, Mode := E_Mode.MAINT_N2, PowerContactorEngaged := TRUE, CablePosM1 := encoderM1.Measurement.CablePosM, CablePosM2 := encoderM2.Measurement.CablePosM, HomedM1 := encoderM1.Homed, HomedM2 := encoderM2.Homed, HomedAndReliableM1 := encoderM1.HomedAndReliable, HomedAndReliableM2 := encoderM2.HomedAndReliable, HomingSuspectM1 := encoderM1.HomingSuspect, HomingSuspectM2 := encoderM2.HomingSuspect, ConfirmClosePosition := btnBucket, Config := cfgBucket, BucketState := bucketState); bucketState := bucket.BucketState;
home.M1Status.HomedAndReliable := encoderM1.HomedAndReliable; home.M2Status.HomedAndReliable := encoderM2.HomedAndReliable; home(BucketOffsetValid := bucketState.BucketReferenced, BtnValidation := bench.Operator.JoyBtnRaw);
ADVANCE_TIME(10000000);
bench(M1_PresetTriggerCmd := encoderM1.HwOut.PresetTriggerCmd, M1_PresetValueOut := encoderM1.HwOut.PresetValueOut, M2_PresetTriggerCmd := encoderM2.HwOut.PresetTriggerCmd, M2_PresetValueOut := encoderM2.HwOut.PresetValueOut, RawPosM1 := raw1, RawPosM2 := raw2); raw1 := bench.RawPosM1; raw2 := bench.RawPosM2;
hw1.RawPosIn := bench.Winch.COD1_PosValue; hw1.SlaveOperational := TRUE; hw2.RawPosIn := bench.Winch.COD2_PosValue; hw2.SlaveOperational := TRUE;
encoderM1(Enable := TRUE, HomingPermit := TRUE, HomingAtTargetM := btnM1, CfgHomingTargetM := 8.7, CfgTopSensorPosM := 8.7, HwIn := hw1, Cfg := cfgEncoder, Calib := calibM1); calibM1 := encoderM1.Calib;
bucketEdge(CLK := btnBucket);
encoderM2(Enable := TRUE, HomingPermit := TRUE, HomingAtTargetM := btnM2 OR bucketEdge.Q, CfgHomingTargetM := 23.7, CfgTopSensorPosM := 23.7, UseDynamicTarget := bucketEdge.Q, DynamicHomingTargetM := encoderM1.Measurement.CablePosM + cfgBucket.OffsetCloseM, HwIn := hw2, Cfg := cfgEncoder, Calib := calibM2); calibM2 := encoderM2.Calib;
bucket(Enable := TRUE, Mode := E_Mode.MAINT_N2, PowerContactorEngaged := TRUE, CablePosM1 := encoderM1.Measurement.CablePosM, CablePosM2 := encoderM2.Measurement.CablePosM, HomedM1 := encoderM1.Homed, HomedM2 := encoderM2.Homed, HomedAndReliableM1 := encoderM1.HomedAndReliable, HomedAndReliableM2 := encoderM2.HomedAndReliable, HomingSuspectM1 := encoderM1.HomingSuspect, HomingSuspectM2 := encoderM2.HomingSuspect, ConfirmClosePosition := btnBucket, Config := cfgBucket, BucketState := bucketState); bucketState := bucket.BucketState;
home.M1Status.HomedAndReliable := encoderM1.HomedAndReliable; home.M2Status.HomedAndReliable := encoderM2.HomedAndReliable; home(BucketOffsetValid := bucketState.BucketReferenced, BtnValidation := bench.Operator.JoyBtnRaw);
ADVANCE_TIME(10000000);
bench(M1_PresetTriggerCmd := encoderM1.HwOut.PresetTriggerCmd, M1_PresetValueOut := encoderM1.HwOut.PresetValueOut, M2_PresetTriggerCmd := encoderM2.HwOut.PresetTriggerCmd, M2_PresetValueOut := encoderM2.HwOut.PresetValueOut, RawPosM1 := raw1, RawPosM2 := raw2); raw1 := bench.RawPosM1; raw2 := bench.RawPosM2;
hw1.RawPosIn := bench.Winch.COD1_PosValue; hw1.SlaveOperational := TRUE; hw2.RawPosIn := bench.Winch.COD2_PosValue; hw2.SlaveOperational := TRUE;
encoderM1(Enable := TRUE, HomingPermit := TRUE, HomingAtTargetM := btnM1, CfgHomingTargetM := 8.7, CfgTopSensorPosM := 8.7, HwIn := hw1, Cfg := cfgEncoder, Calib := calibM1); calibM1 := encoderM1.Calib;
bucketEdge(CLK := btnBucket);
encoderM2(Enable := TRUE, HomingPermit := TRUE, HomingAtTargetM := btnM2 OR bucketEdge.Q, CfgHomingTargetM := 23.7, CfgTopSensorPosM := 23.7, UseDynamicTarget := bucketEdge.Q, DynamicHomingTargetM := encoderM1.Measurement.CablePosM + cfgBucket.OffsetCloseM, HwIn := hw2, Cfg := cfgEncoder, Calib := calibM2); calibM2 := encoderM2.Calib;
bucket(Enable := TRUE, Mode := E_Mode.MAINT_N2, PowerContactorEngaged := TRUE, CablePosM1 := encoderM1.Measurement.CablePosM, CablePosM2 := encoderM2.Measurement.CablePosM, HomedM1 := encoderM1.Homed, HomedM2 := encoderM2.Homed, HomedAndReliableM1 := encoderM1.HomedAndReliable, HomedAndReliableM2 := encoderM2.HomedAndReliable, HomingSuspectM1 := encoderM1.HomingSuspect, HomingSuspectM2 := encoderM2.HomingSuspect, ConfirmClosePosition := btnBucket, Config := cfgBucket, BucketState := bucketState); bucketState := bucket.BucketState;
home.M1Status.HomedAndReliable := encoderM1.HomedAndReliable; home.M2Status.HomedAndReliable := encoderM2.HomedAndReliable; home(BucketOffsetValid := bucketState.BucketReferenced, BtnValidation := bench.Operator.JoyBtnRaw);
ADVANCE_TIME(10000000);
bench(M1_PresetTriggerCmd := encoderM1.HwOut.PresetTriggerCmd, M1_PresetValueOut := encoderM1.HwOut.PresetValueOut, M2_PresetTriggerCmd := encoderM2.HwOut.PresetTriggerCmd, M2_PresetValueOut := encoderM2.HwOut.PresetValueOut, RawPosM1 := raw1, RawPosM2 := raw2); raw1 := bench.RawPosM1; raw2 := bench.RawPosM2;
hw1.RawPosIn := bench.Winch.COD1_PosValue; hw1.SlaveOperational := TRUE; hw2.RawPosIn := bench.Winch.COD2_PosValue; hw2.SlaveOperational := TRUE;
encoderM1(Enable := TRUE, HomingPermit := TRUE, HomingAtTargetM := btnM1, CfgHomingTargetM := 8.7, CfgTopSensorPosM := 8.7, HwIn := hw1, Cfg := cfgEncoder, Calib := calibM1); calibM1 := encoderM1.Calib;
bucketEdge(CLK := btnBucket);
encoderM2(Enable := TRUE, HomingPermit := TRUE, HomingAtTargetM := btnM2 OR bucketEdge.Q, CfgHomingTargetM := 23.7, CfgTopSensorPosM := 23.7, UseDynamicTarget := bucketEdge.Q, DynamicHomingTargetM := encoderM1.Measurement.CablePosM + cfgBucket.OffsetCloseM, HwIn := hw2, Cfg := cfgEncoder, Calib := calibM2); calibM2 := encoderM2.Calib;
bucket(Enable := TRUE, Mode := E_Mode.MAINT_N2, PowerContactorEngaged := TRUE, CablePosM1 := encoderM1.Measurement.CablePosM, CablePosM2 := encoderM2.Measurement.CablePosM, HomedM1 := encoderM1.Homed, HomedM2 := encoderM2.Homed, HomedAndReliableM1 := encoderM1.HomedAndReliable, HomedAndReliableM2 := encoderM2.HomedAndReliable, HomingSuspectM1 := encoderM1.HomingSuspect, HomingSuspectM2 := encoderM2.HomingSuspect, ConfirmClosePosition := btnBucket, Config := cfgBucket, BucketState := bucketState); bucketState := bucket.BucketState;
home.M1Status.HomedAndReliable := encoderM1.HomedAndReliable; home.M2Status.HomedAndReliable := encoderM2.HomedAndReliable; home(BucketOffsetValid := bucketState.BucketReferenced, BtnValidation := bench.Operator.JoyBtnRaw);
ADVANCE_TIME(10000000);
bench(M1_PresetTriggerCmd := encoderM1.HwOut.PresetTriggerCmd, M1_PresetValueOut := encoderM1.HwOut.PresetValueOut, M2_PresetTriggerCmd := encoderM2.HwOut.PresetTriggerCmd, M2_PresetValueOut := encoderM2.HwOut.PresetValueOut, RawPosM1 := raw1, RawPosM2 := raw2); raw1 := bench.RawPosM1; raw2 := bench.RawPosM2;
hw1.RawPosIn := bench.Winch.COD1_PosValue; hw1.SlaveOperational := TRUE; hw2.RawPosIn := bench.Winch.COD2_PosValue; hw2.SlaveOperational := TRUE;
encoderM1(Enable := TRUE, HomingPermit := TRUE, HomingAtTargetM := btnM1, CfgHomingTargetM := 8.7, CfgTopSensorPosM := 8.7, HwIn := hw1, Cfg := cfgEncoder, Calib := calibM1); calibM1 := encoderM1.Calib;
bucketEdge(CLK := btnBucket);
encoderM2(Enable := TRUE, HomingPermit := TRUE, HomingAtTargetM := btnM2 OR bucketEdge.Q, CfgHomingTargetM := 23.7, CfgTopSensorPosM := 23.7, UseDynamicTarget := bucketEdge.Q, DynamicHomingTargetM := encoderM1.Measurement.CablePosM + cfgBucket.OffsetCloseM, HwIn := hw2, Cfg := cfgEncoder, Calib := calibM2); calibM2 := encoderM2.Calib;
bucket(Enable := TRUE, Mode := E_Mode.MAINT_N2, PowerContactorEngaged := TRUE, CablePosM1 := encoderM1.Measurement.CablePosM, CablePosM2 := encoderM2.Measurement.CablePosM, HomedM1 := encoderM1.Homed, HomedM2 := encoderM2.Homed, HomedAndReliableM1 := encoderM1.HomedAndReliable, HomedAndReliableM2 := encoderM2.HomedAndReliable, HomingSuspectM1 := encoderM1.HomingSuspect, HomingSuspectM2 := encoderM2.HomingSuspect, ConfirmClosePosition := btnBucket, Config := cfgBucket, BucketState := bucketState); bucketState := bucket.BucketState;
home.M1Status.HomedAndReliable := encoderM1.HomedAndReliable; home.M2Status.HomedAndReliable := encoderM2.HomedAndReliable; home(BucketOffsetValid := bucketState.BucketReferenced, BtnValidation := bench.Operator.JoyBtnRaw);
ADVANCE_TIME(10000000);
bench(M1_PresetTriggerCmd := encoderM1.HwOut.PresetTriggerCmd, M1_PresetValueOut := encoderM1.HwOut.PresetValueOut, M2_PresetTriggerCmd := encoderM2.HwOut.PresetTriggerCmd, M2_PresetValueOut := encoderM2.HwOut.PresetValueOut, RawPosM1 := raw1, RawPosM2 := raw2); raw1 := bench.RawPosM1; raw2 := bench.RawPosM2;
hw1.RawPosIn := bench.Winch.COD1_PosValue; hw1.SlaveOperational := TRUE; hw2.RawPosIn := bench.Winch.COD2_PosValue; hw2.SlaveOperational := TRUE;
encoderM1(Enable := TRUE, HomingPermit := TRUE, HomingAtTargetM := btnM1, CfgHomingTargetM := 8.7, CfgTopSensorPosM := 8.7, HwIn := hw1, Cfg := cfgEncoder, Calib := calibM1); calibM1 := encoderM1.Calib;
bucketEdge(CLK := btnBucket);
encoderM2(Enable := TRUE, HomingPermit := TRUE, HomingAtTargetM := btnM2 OR bucketEdge.Q, CfgHomingTargetM := 23.7, CfgTopSensorPosM := 23.7, UseDynamicTarget := bucketEdge.Q, DynamicHomingTargetM := encoderM1.Measurement.CablePosM + cfgBucket.OffsetCloseM, HwIn := hw2, Cfg := cfgEncoder, Calib := calibM2); calibM2 := encoderM2.Calib;
bucket(Enable := TRUE, Mode := E_Mode.MAINT_N2, PowerContactorEngaged := TRUE, CablePosM1 := encoderM1.Measurement.CablePosM, CablePosM2 := encoderM2.Measurement.CablePosM, HomedM1 := encoderM1.Homed, HomedM2 := encoderM2.Homed, HomedAndReliableM1 := encoderM1.HomedAndReliable, HomedAndReliableM2 := encoderM2.HomedAndReliable, HomingSuspectM1 := encoderM1.HomingSuspect, HomingSuspectM2 := encoderM2.HomingSuspect, ConfirmClosePosition := btnBucket, Config := cfgBucket, BucketState := bucketState); bucketState := bucket.BucketState;
home.M1Status.HomedAndReliable := encoderM1.HomedAndReliable; home.M2Status.HomedAndReliable := encoderM2.HomedAndReliable; home(BucketOffsetValid := bucketState.BucketReferenced, BtnValidation := bench.Operator.JoyBtnRaw);
ADVANCE_TIME(10000000);
bench(M1_PresetTriggerCmd := encoderM1.HwOut.PresetTriggerCmd, M1_PresetValueOut := encoderM1.HwOut.PresetValueOut, M2_PresetTriggerCmd := encoderM2.HwOut.PresetTriggerCmd, M2_PresetValueOut := encoderM2.HwOut.PresetValueOut, RawPosM1 := raw1, RawPosM2 := raw2); raw1 := bench.RawPosM1; raw2 := bench.RawPosM2;
hw1.RawPosIn := bench.Winch.COD1_PosValue; hw1.SlaveOperational := TRUE; hw2.RawPosIn := bench.Winch.COD2_PosValue; hw2.SlaveOperational := TRUE;
encoderM1(Enable := TRUE, HomingPermit := TRUE, HomingAtTargetM := btnM1, CfgHomingTargetM := 8.7, CfgTopSensorPosM := 8.7, HwIn := hw1, Cfg := cfgEncoder, Calib := calibM1); calibM1 := encoderM1.Calib;
bucketEdge(CLK := btnBucket);
encoderM2(Enable := TRUE, HomingPermit := TRUE, HomingAtTargetM := btnM2 OR bucketEdge.Q, CfgHomingTargetM := 23.7, CfgTopSensorPosM := 23.7, UseDynamicTarget := bucketEdge.Q, DynamicHomingTargetM := encoderM1.Measurement.CablePosM + cfgBucket.OffsetCloseM, HwIn := hw2, Cfg := cfgEncoder, Calib := calibM2); calibM2 := encoderM2.Calib;
bucket(Enable := TRUE, Mode := E_Mode.MAINT_N2, PowerContactorEngaged := TRUE, CablePosM1 := encoderM1.Measurement.CablePosM, CablePosM2 := encoderM2.Measurement.CablePosM, HomedM1 := encoderM1.Homed, HomedM2 := encoderM2.Homed, HomedAndReliableM1 := encoderM1.HomedAndReliable, HomedAndReliableM2 := encoderM2.HomedAndReliable, HomingSuspectM1 := encoderM1.HomingSuspect, HomingSuspectM2 := encoderM2.HomingSuspect, ConfirmClosePosition := btnBucket, Config := cfgBucket, BucketState := bucketState); bucketState := bucket.BucketState;
home.M1Status.HomedAndReliable := encoderM1.HomedAndReliable; home.M2Status.HomedAndReliable := encoderM2.HomedAndReliable; home(BucketOffsetValid := bucketState.BucketReferenced, BtnValidation := bench.Operator.JoyBtnRaw);
ADVANCE_TIME(10000000);
bench(M1_PresetTriggerCmd := encoderM1.HwOut.PresetTriggerCmd, M1_PresetValueOut := encoderM1.HwOut.PresetValueOut, M2_PresetTriggerCmd := encoderM2.HwOut.PresetTriggerCmd, M2_PresetValueOut := encoderM2.HwOut.PresetValueOut, RawPosM1 := raw1, RawPosM2 := raw2); raw1 := bench.RawPosM1; raw2 := bench.RawPosM2;
hw1.RawPosIn := bench.Winch.COD1_PosValue; hw1.SlaveOperational := TRUE; hw2.RawPosIn := bench.Winch.COD2_PosValue; hw2.SlaveOperational := TRUE;
encoderM1(Enable := TRUE, HomingPermit := TRUE, HomingAtTargetM := btnM1, CfgHomingTargetM := 8.7, CfgTopSensorPosM := 8.7, HwIn := hw1, Cfg := cfgEncoder, Calib := calibM1); calibM1 := encoderM1.Calib;
bucketEdge(CLK := btnBucket);
encoderM2(Enable := TRUE, HomingPermit := TRUE, HomingAtTargetM := btnM2 OR bucketEdge.Q, CfgHomingTargetM := 23.7, CfgTopSensorPosM := 23.7, UseDynamicTarget := bucketEdge.Q, DynamicHomingTargetM := encoderM1.Measurement.CablePosM + cfgBucket.OffsetCloseM, HwIn := hw2, Cfg := cfgEncoder, Calib := calibM2); calibM2 := encoderM2.Calib;
bucket(Enable := TRUE, Mode := E_Mode.MAINT_N2, PowerContactorEngaged := TRUE, CablePosM1 := encoderM1.Measurement.CablePosM, CablePosM2 := encoderM2.Measurement.CablePosM, HomedM1 := encoderM1.Homed, HomedM2 := encoderM2.Homed, HomedAndReliableM1 := encoderM1.HomedAndReliable, HomedAndReliableM2 := encoderM2.HomedAndReliable, HomingSuspectM1 := encoderM1.HomingSuspect, HomingSuspectM2 := encoderM2.HomingSuspect, ConfirmClosePosition := btnBucket, Config := cfgBucket, BucketState := bucketState); bucketState := bucket.BucketState;
home.M1Status.HomedAndReliable := encoderM1.HomedAndReliable; home.M2Status.HomedAndReliable := encoderM2.HomedAndReliable; home(BucketOffsetValid := bucketState.BucketReferenced, BtnValidation := bench.Operator.JoyBtnRaw);
ADVANCE_TIME(10000000);
bench(M1_PresetTriggerCmd := encoderM1.HwOut.PresetTriggerCmd, M1_PresetValueOut := encoderM1.HwOut.PresetValueOut, M2_PresetTriggerCmd := encoderM2.HwOut.PresetTriggerCmd, M2_PresetValueOut := encoderM2.HwOut.PresetValueOut, RawPosM1 := raw1, RawPosM2 := raw2); raw1 := bench.RawPosM1; raw2 := bench.RawPosM2;
hw1.RawPosIn := bench.Winch.COD1_PosValue; hw1.SlaveOperational := TRUE; hw2.RawPosIn := bench.Winch.COD2_PosValue; hw2.SlaveOperational := TRUE;
encoderM1(Enable := TRUE, HomingPermit := TRUE, HomingAtTargetM := btnM1, CfgHomingTargetM := 8.7, CfgTopSensorPosM := 8.7, HwIn := hw1, Cfg := cfgEncoder, Calib := calibM1); calibM1 := encoderM1.Calib;
bucketEdge(CLK := btnBucket);
encoderM2(Enable := TRUE, HomingPermit := TRUE, HomingAtTargetM := btnM2 OR bucketEdge.Q, CfgHomingTargetM := 23.7, CfgTopSensorPosM := 23.7, UseDynamicTarget := bucketEdge.Q, DynamicHomingTargetM := encoderM1.Measurement.CablePosM + cfgBucket.OffsetCloseM, HwIn := hw2, Cfg := cfgEncoder, Calib := calibM2); calibM2 := encoderM2.Calib;
bucket(Enable := TRUE, Mode := E_Mode.MAINT_N2, PowerContactorEngaged := TRUE, CablePosM1 := encoderM1.Measurement.CablePosM, CablePosM2 := encoderM2.Measurement.CablePosM, HomedM1 := encoderM1.Homed, HomedM2 := encoderM2.Homed, HomedAndReliableM1 := encoderM1.HomedAndReliable, HomedAndReliableM2 := encoderM2.HomedAndReliable, HomingSuspectM1 := encoderM1.HomingSuspect, HomingSuspectM2 := encoderM2.HomingSuspect, ConfirmClosePosition := btnBucket, Config := cfgBucket, BucketState := bucketState); bucketState := bucket.BucketState;
home.M1Status.HomedAndReliable := encoderM1.HomedAndReliable; home.M2Status.HomedAndReliable := encoderM2.HomedAndReliable; home(BucketOffsetValid := bucketState.BucketReferenced, BtnValidation := bench.Operator.JoyBtnRaw);
ADVANCE_TIME(10000000);
bench(M1_PresetTriggerCmd := encoderM1.HwOut.PresetTriggerCmd, M1_PresetValueOut := encoderM1.HwOut.PresetValueOut, M2_PresetTriggerCmd := encoderM2.HwOut.PresetTriggerCmd, M2_PresetValueOut := encoderM2.HwOut.PresetValueOut, RawPosM1 := raw1, RawPosM2 := raw2); raw1 := bench.RawPosM1; raw2 := bench.RawPosM2;
hw1.RawPosIn := bench.Winch.COD1_PosValue; hw1.SlaveOperational := TRUE; hw2.RawPosIn := bench.Winch.COD2_PosValue; hw2.SlaveOperational := TRUE;
encoderM1(Enable := TRUE, HomingPermit := TRUE, HomingAtTargetM := btnM1, CfgHomingTargetM := 8.7, CfgTopSensorPosM := 8.7, HwIn := hw1, Cfg := cfgEncoder, Calib := calibM1); calibM1 := encoderM1.Calib;
bucketEdge(CLK := btnBucket);
encoderM2(Enable := TRUE, HomingPermit := TRUE, HomingAtTargetM := btnM2 OR bucketEdge.Q, CfgHomingTargetM := 23.7, CfgTopSensorPosM := 23.7, UseDynamicTarget := bucketEdge.Q, DynamicHomingTargetM := encoderM1.Measurement.CablePosM + cfgBucket.OffsetCloseM, HwIn := hw2, Cfg := cfgEncoder, Calib := calibM2); calibM2 := encoderM2.Calib;
bucket(Enable := TRUE, Mode := E_Mode.MAINT_N2, PowerContactorEngaged := TRUE, CablePosM1 := encoderM1.Measurement.CablePosM, CablePosM2 := encoderM2.Measurement.CablePosM, HomedM1 := encoderM1.Homed, HomedM2 := encoderM2.Homed, HomedAndReliableM1 := encoderM1.HomedAndReliable, HomedAndReliableM2 := encoderM2.HomedAndReliable, HomingSuspectM1 := encoderM1.HomingSuspect, HomingSuspectM2 := encoderM2.HomingSuspect, ConfirmClosePosition := btnBucket, Config := cfgBucket, BucketState := bucketState); bucketState := bucket.BucketState;
home.M1Status.HomedAndReliable := encoderM1.HomedAndReliable; home.M2Status.HomedAndReliable := encoderM2.HomedAndReliable; home(BucketOffsetValid := bucketState.BucketReferenced, BtnValidation := bench.Operator.JoyBtnRaw);
ADVANCE_TIME(10000000);
bench(M1_PresetTriggerCmd := encoderM1.HwOut.PresetTriggerCmd, M1_PresetValueOut := encoderM1.HwOut.PresetValueOut, M2_PresetTriggerCmd := encoderM2.HwOut.PresetTriggerCmd, M2_PresetValueOut := encoderM2.HwOut.PresetValueOut, RawPosM1 := raw1, RawPosM2 := raw2); raw1 := bench.RawPosM1; raw2 := bench.RawPosM2;
hw1.RawPosIn := bench.Winch.COD1_PosValue; hw1.SlaveOperational := TRUE; hw2.RawPosIn := bench.Winch.COD2_PosValue; hw2.SlaveOperational := TRUE;
encoderM1(Enable := TRUE, HomingPermit := TRUE, HomingAtTargetM := btnM1, CfgHomingTargetM := 8.7, CfgTopSensorPosM := 8.7, HwIn := hw1, Cfg := cfgEncoder, Calib := calibM1); calibM1 := encoderM1.Calib;
bucketEdge(CLK := btnBucket);
encoderM2(Enable := TRUE, HomingPermit := TRUE, HomingAtTargetM := btnM2 OR bucketEdge.Q, CfgHomingTargetM := 23.7, CfgTopSensorPosM := 23.7, UseDynamicTarget := bucketEdge.Q, DynamicHomingTargetM := encoderM1.Measurement.CablePosM + cfgBucket.OffsetCloseM, HwIn := hw2, Cfg := cfgEncoder, Calib := calibM2); calibM2 := encoderM2.Calib;
bucket(Enable := TRUE, Mode := E_Mode.MAINT_N2, PowerContactorEngaged := TRUE, CablePosM1 := encoderM1.Measurement.CablePosM, CablePosM2 := encoderM2.Measurement.CablePosM, HomedM1 := encoderM1.Homed, HomedM2 := encoderM2.Homed, HomedAndReliableM1 := encoderM1.HomedAndReliable, HomedAndReliableM2 := encoderM2.HomedAndReliable, HomingSuspectM1 := encoderM1.HomingSuspect, HomingSuspectM2 := encoderM2.HomingSuspect, ConfirmClosePosition := btnBucket, Config := cfgBucket, BucketState := bucketState); bucketState := bucket.BucketState;
home.M1Status.HomedAndReliable := encoderM1.HomedAndReliable; home.M2Status.HomedAndReliable := encoderM2.HomedAndReliable; home(BucketOffsetValid := bucketState.BucketReferenced, BtnValidation := bench.Operator.JoyBtnRaw);
ADVANCE_TIME(10000000);
bench(M1_PresetTriggerCmd := encoderM1.HwOut.PresetTriggerCmd, M1_PresetValueOut := encoderM1.HwOut.PresetValueOut, M2_PresetTriggerCmd := encoderM2.HwOut.PresetTriggerCmd, M2_PresetValueOut := encoderM2.HwOut.PresetValueOut, RawPosM1 := raw1, RawPosM2 := raw2); raw1 := bench.RawPosM1; raw2 := bench.RawPosM2;
hw1.RawPosIn := bench.Winch.COD1_PosValue; hw1.SlaveOperational := TRUE; hw2.RawPosIn := bench.Winch.COD2_PosValue; hw2.SlaveOperational := TRUE;
encoderM1(Enable := TRUE, HomingPermit := TRUE, HomingAtTargetM := btnM1, CfgHomingTargetM := 8.7, CfgTopSensorPosM := 8.7, HwIn := hw1, Cfg := cfgEncoder, Calib := calibM1); calibM1 := encoderM1.Calib;
bucketEdge(CLK := btnBucket);
encoderM2(Enable := TRUE, HomingPermit := TRUE, HomingAtTargetM := btnM2 OR bucketEdge.Q, CfgHomingTargetM := 23.7, CfgTopSensorPosM := 23.7, UseDynamicTarget := bucketEdge.Q, DynamicHomingTargetM := encoderM1.Measurement.CablePosM + cfgBucket.OffsetCloseM, HwIn := hw2, Cfg := cfgEncoder, Calib := calibM2); calibM2 := encoderM2.Calib;
bucket(Enable := TRUE, Mode := E_Mode.MAINT_N2, PowerContactorEngaged := TRUE, CablePosM1 := encoderM1.Measurement.CablePosM, CablePosM2 := encoderM2.Measurement.CablePosM, HomedM1 := encoderM1.Homed, HomedM2 := encoderM2.Homed, HomedAndReliableM1 := encoderM1.HomedAndReliable, HomedAndReliableM2 := encoderM2.HomedAndReliable, HomingSuspectM1 := encoderM1.HomingSuspect, HomingSuspectM2 := encoderM2.HomingSuspect, ConfirmClosePosition := btnBucket, Config := cfgBucket, BucketState := bucketState); bucketState := bucket.BucketState;
home.M1Status.HomedAndReliable := encoderM1.HomedAndReliable; home.M2Status.HomedAndReliable := encoderM2.HomedAndReliable; home(BucketOffsetValid := bucketState.BucketReferenced, BtnValidation := bench.Operator.JoyBtnRaw);
ADVANCE_TIME(10000000);
bench(M1_PresetTriggerCmd := encoderM1.HwOut.PresetTriggerCmd, M1_PresetValueOut := encoderM1.HwOut.PresetValueOut, M2_PresetTriggerCmd := encoderM2.HwOut.PresetTriggerCmd, M2_PresetValueOut := encoderM2.HwOut.PresetValueOut, RawPosM1 := raw1, RawPosM2 := raw2); raw1 := bench.RawPosM1; raw2 := bench.RawPosM2;
hw1.RawPosIn := bench.Winch.COD1_PosValue; hw1.SlaveOperational := TRUE; hw2.RawPosIn := bench.Winch.COD2_PosValue; hw2.SlaveOperational := TRUE;
encoderM1(Enable := TRUE, HomingPermit := TRUE, HomingAtTargetM := btnM1, CfgHomingTargetM := 8.7, CfgTopSensorPosM := 8.7, HwIn := hw1, Cfg := cfgEncoder, Calib := calibM1); calibM1 := encoderM1.Calib;
bucketEdge(CLK := btnBucket);
encoderM2(Enable := TRUE, HomingPermit := TRUE, HomingAtTargetM := btnM2 OR bucketEdge.Q, CfgHomingTargetM := 23.7, CfgTopSensorPosM := 23.7, UseDynamicTarget := bucketEdge.Q, DynamicHomingTargetM := encoderM1.Measurement.CablePosM + cfgBucket.OffsetCloseM, HwIn := hw2, Cfg := cfgEncoder, Calib := calibM2); calibM2 := encoderM2.Calib;
bucket(Enable := TRUE, Mode := E_Mode.MAINT_N2, PowerContactorEngaged := TRUE, CablePosM1 := encoderM1.Measurement.CablePosM, CablePosM2 := encoderM2.Measurement.CablePosM, HomedM1 := encoderM1.Homed, HomedM2 := encoderM2.Homed, HomedAndReliableM1 := encoderM1.HomedAndReliable, HomedAndReliableM2 := encoderM2.HomedAndReliable, HomingSuspectM1 := encoderM1.HomingSuspect, HomingSuspectM2 := encoderM2.HomingSuspect, ConfirmClosePosition := btnBucket, Config := cfgBucket, BucketState := bucketState); bucketState := bucket.BucketState;
home.M1Status.HomedAndReliable := encoderM1.HomedAndReliable; home.M2Status.HomedAndReliable := encoderM2.HomedAndReliable; home(BucketOffsetValid := bucketState.BucketReferenced, BtnValidation := bench.Operator.JoyBtnRaw);
ADVANCE_TIME(10000000);
bench(M1_PresetTriggerCmd := encoderM1.HwOut.PresetTriggerCmd, M1_PresetValueOut := encoderM1.HwOut.PresetValueOut, M2_PresetTriggerCmd := encoderM2.HwOut.PresetTriggerCmd, M2_PresetValueOut := encoderM2.HwOut.PresetValueOut, RawPosM1 := raw1, RawPosM2 := raw2); raw1 := bench.RawPosM1; raw2 := bench.RawPosM2;
hw1.RawPosIn := bench.Winch.COD1_PosValue; hw1.SlaveOperational := TRUE; hw2.RawPosIn := bench.Winch.COD2_PosValue; hw2.SlaveOperational := TRUE;
encoderM1(Enable := TRUE, HomingPermit := TRUE, HomingAtTargetM := btnM1, CfgHomingTargetM := 8.7, CfgTopSensorPosM := 8.7, HwIn := hw1, Cfg := cfgEncoder, Calib := calibM1); calibM1 := encoderM1.Calib;
bucketEdge(CLK := btnBucket);
encoderM2(Enable := TRUE, HomingPermit := TRUE, HomingAtTargetM := btnM2 OR bucketEdge.Q, CfgHomingTargetM := 23.7, CfgTopSensorPosM := 23.7, UseDynamicTarget := bucketEdge.Q, DynamicHomingTargetM := encoderM1.Measurement.CablePosM + cfgBucket.OffsetCloseM, HwIn := hw2, Cfg := cfgEncoder, Calib := calibM2); calibM2 := encoderM2.Calib;
bucket(Enable := TRUE, Mode := E_Mode.MAINT_N2, PowerContactorEngaged := TRUE, CablePosM1 := encoderM1.Measurement.CablePosM, CablePosM2 := encoderM2.Measurement.CablePosM, HomedM1 := encoderM1.Homed, HomedM2 := encoderM2.Homed, HomedAndReliableM1 := encoderM1.HomedAndReliable, HomedAndReliableM2 := encoderM2.HomedAndReliable, HomingSuspectM1 := encoderM1.HomingSuspect, HomingSuspectM2 := encoderM2.HomingSuspect, ConfirmClosePosition := btnBucket, Config := cfgBucket, BucketState := bucketState); bucketState := bucket.BucketState;
home.M1Status.HomedAndReliable := encoderM1.HomedAndReliable; home.M2Status.HomedAndReliable := encoderM2.HomedAndReliable; home(BucketOffsetValid := bucketState.BucketReferenced, BtnValidation := bench.Operator.JoyBtnRaw);
ADVANCE_TIME(10000000);
bench(M1_PresetTriggerCmd := encoderM1.HwOut.PresetTriggerCmd, M1_PresetValueOut := encoderM1.HwOut.PresetValueOut, M2_PresetTriggerCmd := encoderM2.HwOut.PresetTriggerCmd, M2_PresetValueOut := encoderM2.HwOut.PresetValueOut, RawPosM1 := raw1, RawPosM2 := raw2); raw1 := bench.RawPosM1; raw2 := bench.RawPosM2;
hw1.RawPosIn := bench.Winch.COD1_PosValue; hw1.SlaveOperational := TRUE; hw2.RawPosIn := bench.Winch.COD2_PosValue; hw2.SlaveOperational := TRUE;
encoderM1(Enable := TRUE, HomingPermit := TRUE, HomingAtTargetM := btnM1, CfgHomingTargetM := 8.7, CfgTopSensorPosM := 8.7, HwIn := hw1, Cfg := cfgEncoder, Calib := calibM1); calibM1 := encoderM1.Calib;
bucketEdge(CLK := btnBucket);
encoderM2(Enable := TRUE, HomingPermit := TRUE, HomingAtTargetM := btnM2 OR bucketEdge.Q, CfgHomingTargetM := 23.7, CfgTopSensorPosM := 23.7, UseDynamicTarget := bucketEdge.Q, DynamicHomingTargetM := encoderM1.Measurement.CablePosM + cfgBucket.OffsetCloseM, HwIn := hw2, Cfg := cfgEncoder, Calib := calibM2); calibM2 := encoderM2.Calib;
bucket(Enable := TRUE, Mode := E_Mode.MAINT_N2, PowerContactorEngaged := TRUE, CablePosM1 := encoderM1.Measurement.CablePosM, CablePosM2 := encoderM2.Measurement.CablePosM, HomedM1 := encoderM1.Homed, HomedM2 := encoderM2.Homed, HomedAndReliableM1 := encoderM1.HomedAndReliable, HomedAndReliableM2 := encoderM2.HomedAndReliable, HomingSuspectM1 := encoderM1.HomingSuspect, HomingSuspectM2 := encoderM2.HomingSuspect, ConfirmClosePosition := btnBucket, Config := cfgBucket, BucketState := bucketState); bucketState := bucket.BucketState;
home.M1Status.HomedAndReliable := encoderM1.HomedAndReliable; home.M2Status.HomedAndReliable := encoderM2.HomedAndReliable; home(BucketOffsetValid := bucketState.BucketReferenced, BtnValidation := bench.Operator.JoyBtnRaw);
ADVANCE_TIME(10000000);
bench(M1_PresetTriggerCmd := encoderM1.HwOut.PresetTriggerCmd, M1_PresetValueOut := encoderM1.HwOut.PresetValueOut, M2_PresetTriggerCmd := encoderM2.HwOut.PresetTriggerCmd, M2_PresetValueOut := encoderM2.HwOut.PresetValueOut, RawPosM1 := raw1, RawPosM2 := raw2); raw1 := bench.RawPosM1; raw2 := bench.RawPosM2;
hw1.RawPosIn := bench.Winch.COD1_PosValue; hw1.SlaveOperational := TRUE; hw2.RawPosIn := bench.Winch.COD2_PosValue; hw2.SlaveOperational := TRUE;
encoderM1(Enable := TRUE, HomingPermit := TRUE, HomingAtTargetM := btnM1, CfgHomingTargetM := 8.7, CfgTopSensorPosM := 8.7, HwIn := hw1, Cfg := cfgEncoder, Calib := calibM1); calibM1 := encoderM1.Calib;
bucketEdge(CLK := btnBucket);
encoderM2(Enable := TRUE, HomingPermit := TRUE, HomingAtTargetM := btnM2 OR bucketEdge.Q, CfgHomingTargetM := 23.7, CfgTopSensorPosM := 23.7, UseDynamicTarget := bucketEdge.Q, DynamicHomingTargetM := encoderM1.Measurement.CablePosM + cfgBucket.OffsetCloseM, HwIn := hw2, Cfg := cfgEncoder, Calib := calibM2); calibM2 := encoderM2.Calib;
bucket(Enable := TRUE, Mode := E_Mode.MAINT_N2, PowerContactorEngaged := TRUE, CablePosM1 := encoderM1.Measurement.CablePosM, CablePosM2 := encoderM2.Measurement.CablePosM, HomedM1 := encoderM1.Homed, HomedM2 := encoderM2.Homed, HomedAndReliableM1 := encoderM1.HomedAndReliable, HomedAndReliableM2 := encoderM2.HomedAndReliable, HomingSuspectM1 := encoderM1.HomingSuspect, HomingSuspectM2 := encoderM2.HomingSuspect, ConfirmClosePosition := btnBucket, Config := cfgBucket, BucketState := bucketState); bucketState := bucket.BucketState;
home.M1Status.HomedAndReliable := encoderM1.HomedAndReliable; home.M2Status.HomedAndReliable := encoderM2.HomedAndReliable; home(BucketOffsetValid := bucketState.BucketReferenced, BtnValidation := bench.Operator.JoyBtnRaw);
ADVANCE_TIME(10000000);
bench(M1_PresetTriggerCmd := encoderM1.HwOut.PresetTriggerCmd, M1_PresetValueOut := encoderM1.HwOut.PresetValueOut, M2_PresetTriggerCmd := encoderM2.HwOut.PresetTriggerCmd, M2_PresetValueOut := encoderM2.HwOut.PresetValueOut, RawPosM1 := raw1, RawPosM2 := raw2); raw1 := bench.RawPosM1; raw2 := bench.RawPosM2;
hw1.RawPosIn := bench.Winch.COD1_PosValue; hw1.SlaveOperational := TRUE; hw2.RawPosIn := bench.Winch.COD2_PosValue; hw2.SlaveOperational := TRUE;
encoderM1(Enable := TRUE, HomingPermit := TRUE, HomingAtTargetM := btnM1, CfgHomingTargetM := 8.7, CfgTopSensorPosM := 8.7, HwIn := hw1, Cfg := cfgEncoder, Calib := calibM1); calibM1 := encoderM1.Calib;
bucketEdge(CLK := btnBucket);
encoderM2(Enable := TRUE, HomingPermit := TRUE, HomingAtTargetM := btnM2 OR bucketEdge.Q, CfgHomingTargetM := 23.7, CfgTopSensorPosM := 23.7, UseDynamicTarget := bucketEdge.Q, DynamicHomingTargetM := encoderM1.Measurement.CablePosM + cfgBucket.OffsetCloseM, HwIn := hw2, Cfg := cfgEncoder, Calib := calibM2); calibM2 := encoderM2.Calib;
bucket(Enable := TRUE, Mode := E_Mode.MAINT_N2, PowerContactorEngaged := TRUE, CablePosM1 := encoderM1.Measurement.CablePosM, CablePosM2 := encoderM2.Measurement.CablePosM, HomedM1 := encoderM1.Homed, HomedM2 := encoderM2.Homed, HomedAndReliableM1 := encoderM1.HomedAndReliable, HomedAndReliableM2 := encoderM2.HomedAndReliable, HomingSuspectM1 := encoderM1.HomingSuspect, HomingSuspectM2 := encoderM2.HomingSuspect, ConfirmClosePosition := btnBucket, Config := cfgBucket, BucketState := bucketState); bucketState := bucket.BucketState;
home.M1Status.HomedAndReliable := encoderM1.HomedAndReliable; home.M2Status.HomedAndReliable := encoderM2.HomedAndReliable; home(BucketOffsetValid := bucketState.BucketReferenced, BtnValidation := bench.Operator.JoyBtnRaw);
ADVANCE_TIME(10000000);
bench(M1_PresetTriggerCmd := encoderM1.HwOut.PresetTriggerCmd, M1_PresetValueOut := encoderM1.HwOut.PresetValueOut, M2_PresetTriggerCmd := encoderM2.HwOut.PresetTriggerCmd, M2_PresetValueOut := encoderM2.HwOut.PresetValueOut, RawPosM1 := raw1, RawPosM2 := raw2); raw1 := bench.RawPosM1; raw2 := bench.RawPosM2;
hw1.RawPosIn := bench.Winch.COD1_PosValue; hw1.SlaveOperational := TRUE; hw2.RawPosIn := bench.Winch.COD2_PosValue; hw2.SlaveOperational := TRUE;
encoderM1(Enable := TRUE, HomingPermit := TRUE, HomingAtTargetM := btnM1, CfgHomingTargetM := 8.7, CfgTopSensorPosM := 8.7, HwIn := hw1, Cfg := cfgEncoder, Calib := calibM1); calibM1 := encoderM1.Calib;
bucketEdge(CLK := btnBucket);
encoderM2(Enable := TRUE, HomingPermit := TRUE, HomingAtTargetM := btnM2 OR bucketEdge.Q, CfgHomingTargetM := 23.7, CfgTopSensorPosM := 23.7, UseDynamicTarget := bucketEdge.Q, DynamicHomingTargetM := encoderM1.Measurement.CablePosM + cfgBucket.OffsetCloseM, HwIn := hw2, Cfg := cfgEncoder, Calib := calibM2); calibM2 := encoderM2.Calib;
bucket(Enable := TRUE, Mode := E_Mode.MAINT_N2, PowerContactorEngaged := TRUE, CablePosM1 := encoderM1.Measurement.CablePosM, CablePosM2 := encoderM2.Measurement.CablePosM, HomedM1 := encoderM1.Homed, HomedM2 := encoderM2.Homed, HomedAndReliableM1 := encoderM1.HomedAndReliable, HomedAndReliableM2 := encoderM2.HomedAndReliable, HomingSuspectM1 := encoderM1.HomingSuspect, HomingSuspectM2 := encoderM2.HomingSuspect, ConfirmClosePosition := btnBucket, Config := cfgBucket, BucketState := bucketState); bucketState := bucket.BucketState;
home.M1Status.HomedAndReliable := encoderM1.HomedAndReliable; home.M2Status.HomedAndReliable := encoderM2.HomedAndReliable; home(BucketOffsetValid := bucketState.BucketReferenced, BtnValidation := bench.Operator.JoyBtnRaw);
ADVANCE_TIME(10000000);
bench(M1_PresetTriggerCmd := encoderM1.HwOut.PresetTriggerCmd, M1_PresetValueOut := encoderM1.HwOut.PresetValueOut, M2_PresetTriggerCmd := encoderM2.HwOut.PresetTriggerCmd, M2_PresetValueOut := encoderM2.HwOut.PresetValueOut, RawPosM1 := raw1, RawPosM2 := raw2); raw1 := bench.RawPosM1; raw2 := bench.RawPosM2;
hw1.RawPosIn := bench.Winch.COD1_PosValue; hw1.SlaveOperational := TRUE; hw2.RawPosIn := bench.Winch.COD2_PosValue; hw2.SlaveOperational := TRUE;
encoderM1(Enable := TRUE, HomingPermit := TRUE, HomingAtTargetM := btnM1, CfgHomingTargetM := 8.7, CfgTopSensorPosM := 8.7, HwIn := hw1, Cfg := cfgEncoder, Calib := calibM1); calibM1 := encoderM1.Calib;
bucketEdge(CLK := btnBucket);
encoderM2(Enable := TRUE, HomingPermit := TRUE, HomingAtTargetM := btnM2 OR bucketEdge.Q, CfgHomingTargetM := 23.7, CfgTopSensorPosM := 23.7, UseDynamicTarget := bucketEdge.Q, DynamicHomingTargetM := encoderM1.Measurement.CablePosM + cfgBucket.OffsetCloseM, HwIn := hw2, Cfg := cfgEncoder, Calib := calibM2); calibM2 := encoderM2.Calib;
bucket(Enable := TRUE, Mode := E_Mode.MAINT_N2, PowerContactorEngaged := TRUE, CablePosM1 := encoderM1.Measurement.CablePosM, CablePosM2 := encoderM2.Measurement.CablePosM, HomedM1 := encoderM1.Homed, HomedM2 := encoderM2.Homed, HomedAndReliableM1 := encoderM1.HomedAndReliable, HomedAndReliableM2 := encoderM2.HomedAndReliable, HomingSuspectM1 := encoderM1.HomingSuspect, HomingSuspectM2 := encoderM2.HomingSuspect, ConfirmClosePosition := btnBucket, Config := cfgBucket, BucketState := bucketState); bucketState := bucket.BucketState;
home.M1Status.HomedAndReliable := encoderM1.HomedAndReliable; home.M2Status.HomedAndReliable := encoderM2.HomedAndReliable; home(BucketOffsetValid := bucketState.BucketReferenced, BtnValidation := bench.Operator.JoyBtnRaw);
ADVANCE_TIME(10000000);
bench(M1_PresetTriggerCmd := encoderM1.HwOut.PresetTriggerCmd, M1_PresetValueOut := encoderM1.HwOut.PresetValueOut, M2_PresetTriggerCmd := encoderM2.HwOut.PresetTriggerCmd, M2_PresetValueOut := encoderM2.HwOut.PresetValueOut, RawPosM1 := raw1, RawPosM2 := raw2); raw1 := bench.RawPosM1; raw2 := bench.RawPosM2;
hw1.RawPosIn := bench.Winch.COD1_PosValue; hw1.SlaveOperational := TRUE; hw2.RawPosIn := bench.Winch.COD2_PosValue; hw2.SlaveOperational := TRUE;
encoderM1(Enable := TRUE, HomingPermit := TRUE, HomingAtTargetM := btnM1, CfgHomingTargetM := 8.7, CfgTopSensorPosM := 8.7, HwIn := hw1, Cfg := cfgEncoder, Calib := calibM1); calibM1 := encoderM1.Calib;
bucketEdge(CLK := btnBucket);
encoderM2(Enable := TRUE, HomingPermit := TRUE, HomingAtTargetM := btnM2 OR bucketEdge.Q, CfgHomingTargetM := 23.7, CfgTopSensorPosM := 23.7, UseDynamicTarget := bucketEdge.Q, DynamicHomingTargetM := encoderM1.Measurement.CablePosM + cfgBucket.OffsetCloseM, HwIn := hw2, Cfg := cfgEncoder, Calib := calibM2); calibM2 := encoderM2.Calib;
bucket(Enable := TRUE, Mode := E_Mode.MAINT_N2, PowerContactorEngaged := TRUE, CablePosM1 := encoderM1.Measurement.CablePosM, CablePosM2 := encoderM2.Measurement.CablePosM, HomedM1 := encoderM1.Homed, HomedM2 := encoderM2.Homed, HomedAndReliableM1 := encoderM1.HomedAndReliable, HomedAndReliableM2 := encoderM2.HomedAndReliable, HomingSuspectM1 := encoderM1.HomingSuspect, HomingSuspectM2 := encoderM2.HomingSuspect, ConfirmClosePosition := btnBucket, Config := cfgBucket, BucketState := bucketState); bucketState := bucket.BucketState;
home.M1Status.HomedAndReliable := encoderM1.HomedAndReliable; home.M2Status.HomedAndReliable := encoderM2.HomedAndReliable; home(BucketOffsetValid := bucketState.BucketReferenced, BtnValidation := bench.Operator.JoyBtnRaw);
ADVANCE_TIME(10000000);
bench(M1_PresetTriggerCmd := encoderM1.HwOut.PresetTriggerCmd, M1_PresetValueOut := encoderM1.HwOut.PresetValueOut, M2_PresetTriggerCmd := encoderM2.HwOut.PresetTriggerCmd, M2_PresetValueOut := encoderM2.HwOut.PresetValueOut, RawPosM1 := raw1, RawPosM2 := raw2); raw1 := bench.RawPosM1; raw2 := bench.RawPosM2;
hw1.RawPosIn := bench.Winch.COD1_PosValue; hw1.SlaveOperational := TRUE; hw2.RawPosIn := bench.Winch.COD2_PosValue; hw2.SlaveOperational := TRUE;
encoderM1(Enable := TRUE, HomingPermit := TRUE, HomingAtTargetM := btnM1, CfgHomingTargetM := 8.7, CfgTopSensorPosM := 8.7, HwIn := hw1, Cfg := cfgEncoder, Calib := calibM1); calibM1 := encoderM1.Calib;
bucketEdge(CLK := btnBucket);
encoderM2(Enable := TRUE, HomingPermit := TRUE, HomingAtTargetM := btnM2 OR bucketEdge.Q, CfgHomingTargetM := 23.7, CfgTopSensorPosM := 23.7, UseDynamicTarget := bucketEdge.Q, DynamicHomingTargetM := encoderM1.Measurement.CablePosM + cfgBucket.OffsetCloseM, HwIn := hw2, Cfg := cfgEncoder, Calib := calibM2); calibM2 := encoderM2.Calib;
bucket(Enable := TRUE, Mode := E_Mode.MAINT_N2, PowerContactorEngaged := TRUE, CablePosM1 := encoderM1.Measurement.CablePosM, CablePosM2 := encoderM2.Measurement.CablePosM, HomedM1 := encoderM1.Homed, HomedM2 := encoderM2.Homed, HomedAndReliableM1 := encoderM1.HomedAndReliable, HomedAndReliableM2 := encoderM2.HomedAndReliable, HomingSuspectM1 := encoderM1.HomingSuspect, HomingSuspectM2 := encoderM2.HomingSuspect, ConfirmClosePosition := btnBucket, Config := cfgBucket, BucketState := bucketState); bucketState := bucket.BucketState;
home.M1Status.HomedAndReliable := encoderM1.HomedAndReliable; home.M2Status.HomedAndReliable := encoderM2.HomedAndReliable; home(BucketOffsetValid := bucketState.BucketReferenced, BtnValidation := bench.Operator.JoyBtnRaw);
ADVANCE_TIME(10000000);
bench(M1_PresetTriggerCmd := encoderM1.HwOut.PresetTriggerCmd, M1_PresetValueOut := encoderM1.HwOut.PresetValueOut, M2_PresetTriggerCmd := encoderM2.HwOut.PresetTriggerCmd, M2_PresetValueOut := encoderM2.HwOut.PresetValueOut, RawPosM1 := raw1, RawPosM2 := raw2); raw1 := bench.RawPosM1; raw2 := bench.RawPosM2;
hw1.RawPosIn := bench.Winch.COD1_PosValue; hw1.SlaveOperational := TRUE; hw2.RawPosIn := bench.Winch.COD2_PosValue; hw2.SlaveOperational := TRUE;
encoderM1(Enable := TRUE, HomingPermit := TRUE, HomingAtTargetM := btnM1, CfgHomingTargetM := 8.7, CfgTopSensorPosM := 8.7, HwIn := hw1, Cfg := cfgEncoder, Calib := calibM1); calibM1 := encoderM1.Calib;
bucketEdge(CLK := btnBucket);
encoderM2(Enable := TRUE, HomingPermit := TRUE, HomingAtTargetM := btnM2 OR bucketEdge.Q, CfgHomingTargetM := 23.7, CfgTopSensorPosM := 23.7, UseDynamicTarget := bucketEdge.Q, DynamicHomingTargetM := encoderM1.Measurement.CablePosM + cfgBucket.OffsetCloseM, HwIn := hw2, Cfg := cfgEncoder, Calib := calibM2); calibM2 := encoderM2.Calib;
bucket(Enable := TRUE, Mode := E_Mode.MAINT_N2, PowerContactorEngaged := TRUE, CablePosM1 := encoderM1.Measurement.CablePosM, CablePosM2 := encoderM2.Measurement.CablePosM, HomedM1 := encoderM1.Homed, HomedM2 := encoderM2.Homed, HomedAndReliableM1 := encoderM1.HomedAndReliable, HomedAndReliableM2 := encoderM2.HomedAndReliable, HomingSuspectM1 := encoderM1.HomingSuspect, HomingSuspectM2 := encoderM2.HomingSuspect, ConfirmClosePosition := btnBucket, Config := cfgBucket, BucketState := bucketState); bucketState := bucket.BucketState;
home.M1Status.HomedAndReliable := encoderM1.HomedAndReliable; home.M2Status.HomedAndReliable := encoderM2.HomedAndReliable; home(BucketOffsetValid := bucketState.BucketReferenced, BtnValidation := bench.Operator.JoyBtnRaw);
ADVANCE_TIME(10000000);
bench(M1_PresetTriggerCmd := encoderM1.HwOut.PresetTriggerCmd, M1_PresetValueOut := encoderM1.HwOut.PresetValueOut, M2_PresetTriggerCmd := encoderM2.HwOut.PresetTriggerCmd, M2_PresetValueOut := encoderM2.HwOut.PresetValueOut, RawPosM1 := raw1, RawPosM2 := raw2); raw1 := bench.RawPosM1; raw2 := bench.RawPosM2;
hw1.RawPosIn := bench.Winch.COD1_PosValue; hw1.SlaveOperational := TRUE; hw2.RawPosIn := bench.Winch.COD2_PosValue; hw2.SlaveOperational := TRUE;
encoderM1(Enable := TRUE, HomingPermit := TRUE, HomingAtTargetM := btnM1, CfgHomingTargetM := 8.7, CfgTopSensorPosM := 8.7, HwIn := hw1, Cfg := cfgEncoder, Calib := calibM1); calibM1 := encoderM1.Calib;
bucketEdge(CLK := btnBucket);
encoderM2(Enable := TRUE, HomingPermit := TRUE, HomingAtTargetM := btnM2 OR bucketEdge.Q, CfgHomingTargetM := 23.7, CfgTopSensorPosM := 23.7, UseDynamicTarget := bucketEdge.Q, DynamicHomingTargetM := encoderM1.Measurement.CablePosM + cfgBucket.OffsetCloseM, HwIn := hw2, Cfg := cfgEncoder, Calib := calibM2); calibM2 := encoderM2.Calib;
bucket(Enable := TRUE, Mode := E_Mode.MAINT_N2, PowerContactorEngaged := TRUE, CablePosM1 := encoderM1.Measurement.CablePosM, CablePosM2 := encoderM2.Measurement.CablePosM, HomedM1 := encoderM1.Homed, HomedM2 := encoderM2.Homed, HomedAndReliableM1 := encoderM1.HomedAndReliable, HomedAndReliableM2 := encoderM2.HomedAndReliable, HomingSuspectM1 := encoderM1.HomingSuspect, HomingSuspectM2 := encoderM2.HomingSuspect, ConfirmClosePosition := btnBucket, Config := cfgBucket, BucketState := bucketState); bucketState := bucket.BucketState;
home.M1Status.HomedAndReliable := encoderM1.HomedAndReliable; home.M2Status.HomedAndReliable := encoderM2.HomedAndReliable; home(BucketOffsetValid := bucketState.BucketReferenced, BtnValidation := bench.Operator.JoyBtnRaw);
ADVANCE_TIME(10000000);
bench(M1_PresetTriggerCmd := encoderM1.HwOut.PresetTriggerCmd, M1_PresetValueOut := encoderM1.HwOut.PresetValueOut, M2_PresetTriggerCmd := encoderM2.HwOut.PresetTriggerCmd, M2_PresetValueOut := encoderM2.HwOut.PresetValueOut, RawPosM1 := raw1, RawPosM2 := raw2); raw1 := bench.RawPosM1; raw2 := bench.RawPosM2;
hw1.RawPosIn := bench.Winch.COD1_PosValue; hw1.SlaveOperational := TRUE; hw2.RawPosIn := bench.Winch.COD2_PosValue; hw2.SlaveOperational := TRUE;
encoderM1(Enable := TRUE, HomingPermit := TRUE, HomingAtTargetM := btnM1, CfgHomingTargetM := 8.7, CfgTopSensorPosM := 8.7, HwIn := hw1, Cfg := cfgEncoder, Calib := calibM1); calibM1 := encoderM1.Calib;
bucketEdge(CLK := btnBucket);
encoderM2(Enable := TRUE, HomingPermit := TRUE, HomingAtTargetM := btnM2 OR bucketEdge.Q, CfgHomingTargetM := 23.7, CfgTopSensorPosM := 23.7, UseDynamicTarget := bucketEdge.Q, DynamicHomingTargetM := encoderM1.Measurement.CablePosM + cfgBucket.OffsetCloseM, HwIn := hw2, Cfg := cfgEncoder, Calib := calibM2); calibM2 := encoderM2.Calib;
bucket(Enable := TRUE, Mode := E_Mode.MAINT_N2, PowerContactorEngaged := TRUE, CablePosM1 := encoderM1.Measurement.CablePosM, CablePosM2 := encoderM2.Measurement.CablePosM, HomedM1 := encoderM1.Homed, HomedM2 := encoderM2.Homed, HomedAndReliableM1 := encoderM1.HomedAndReliable, HomedAndReliableM2 := encoderM2.HomedAndReliable, HomingSuspectM1 := encoderM1.HomingSuspect, HomingSuspectM2 := encoderM2.HomingSuspect, ConfirmClosePosition := btnBucket, Config := cfgBucket, BucketState := bucketState); bucketState := bucket.BucketState;
home.M1Status.HomedAndReliable := encoderM1.HomedAndReliable; home.M2Status.HomedAndReliable := encoderM2.HomedAndReliable; home(BucketOffsetValid := bucketState.BucketReferenced, BtnValidation := bench.Operator.JoyBtnRaw);
ADVANCE_TIME(10000000);
bench(M1_PresetTriggerCmd := encoderM1.HwOut.PresetTriggerCmd, M1_PresetValueOut := encoderM1.HwOut.PresetValueOut, M2_PresetTriggerCmd := encoderM2.HwOut.PresetTriggerCmd, M2_PresetValueOut := encoderM2.HwOut.PresetValueOut, RawPosM1 := raw1, RawPosM2 := raw2); raw1 := bench.RawPosM1; raw2 := bench.RawPosM2;
hw1.RawPosIn := bench.Winch.COD1_PosValue; hw1.SlaveOperational := TRUE; hw2.RawPosIn := bench.Winch.COD2_PosValue; hw2.SlaveOperational := TRUE;
encoderM1(Enable := TRUE, HomingPermit := TRUE, HomingAtTargetM := btnM1, CfgHomingTargetM := 8.7, CfgTopSensorPosM := 8.7, HwIn := hw1, Cfg := cfgEncoder, Calib := calibM1); calibM1 := encoderM1.Calib;
bucketEdge(CLK := btnBucket);
encoderM2(Enable := TRUE, HomingPermit := TRUE, HomingAtTargetM := btnM2 OR bucketEdge.Q, CfgHomingTargetM := 23.7, CfgTopSensorPosM := 23.7, UseDynamicTarget := bucketEdge.Q, DynamicHomingTargetM := encoderM1.Measurement.CablePosM + cfgBucket.OffsetCloseM, HwIn := hw2, Cfg := cfgEncoder, Calib := calibM2); calibM2 := encoderM2.Calib;
bucket(Enable := TRUE, Mode := E_Mode.MAINT_N2, PowerContactorEngaged := TRUE, CablePosM1 := encoderM1.Measurement.CablePosM, CablePosM2 := encoderM2.Measurement.CablePosM, HomedM1 := encoderM1.Homed, HomedM2 := encoderM2.Homed, HomedAndReliableM1 := encoderM1.HomedAndReliable, HomedAndReliableM2 := encoderM2.HomedAndReliable, HomingSuspectM1 := encoderM1.HomingSuspect, HomingSuspectM2 := encoderM2.HomingSuspect, ConfirmClosePosition := btnBucket, Config := cfgBucket, BucketState := bucketState); bucketState := bucket.BucketState;
home.M1Status.HomedAndReliable := encoderM1.HomedAndReliable; home.M2Status.HomedAndReliable := encoderM2.HomedAndReliable; home(BucketOffsetValid := bucketState.BucketReferenced, BtnValidation := bench.Operator.JoyBtnRaw);
ADVANCE_TIME(10000000);
bench(M1_PresetTriggerCmd := encoderM1.HwOut.PresetTriggerCmd, M1_PresetValueOut := encoderM1.HwOut.PresetValueOut, M2_PresetTriggerCmd := encoderM2.HwOut.PresetTriggerCmd, M2_PresetValueOut := encoderM2.HwOut.PresetValueOut, RawPosM1 := raw1, RawPosM2 := raw2); raw1 := bench.RawPosM1; raw2 := bench.RawPosM2;
hw1.RawPosIn := bench.Winch.COD1_PosValue; hw1.SlaveOperational := TRUE; hw2.RawPosIn := bench.Winch.COD2_PosValue; hw2.SlaveOperational := TRUE;
encoderM1(Enable := TRUE, HomingPermit := TRUE, HomingAtTargetM := btnM1, CfgHomingTargetM := 8.7, CfgTopSensorPosM := 8.7, HwIn := hw1, Cfg := cfgEncoder, Calib := calibM1); calibM1 := encoderM1.Calib;
bucketEdge(CLK := btnBucket);
encoderM2(Enable := TRUE, HomingPermit := TRUE, HomingAtTargetM := btnM2 OR bucketEdge.Q, CfgHomingTargetM := 23.7, CfgTopSensorPosM := 23.7, UseDynamicTarget := bucketEdge.Q, DynamicHomingTargetM := encoderM1.Measurement.CablePosM + cfgBucket.OffsetCloseM, HwIn := hw2, Cfg := cfgEncoder, Calib := calibM2); calibM2 := encoderM2.Calib;
bucket(Enable := TRUE, Mode := E_Mode.MAINT_N2, PowerContactorEngaged := TRUE, CablePosM1 := encoderM1.Measurement.CablePosM, CablePosM2 := encoderM2.Measurement.CablePosM, HomedM1 := encoderM1.Homed, HomedM2 := encoderM2.Homed, HomedAndReliableM1 := encoderM1.HomedAndReliable, HomedAndReliableM2 := encoderM2.HomedAndReliable, HomingSuspectM1 := encoderM1.HomingSuspect, HomingSuspectM2 := encoderM2.HomingSuspect, ConfirmClosePosition := btnBucket, Config := cfgBucket, BucketState := bucketState); bucketState := bucket.BucketState;
home.M1Status.HomedAndReliable := encoderM1.HomedAndReliable; home.M2Status.HomedAndReliable := encoderM2.HomedAndReliable; home(BucketOffsetValid := bucketState.BucketReferenced, BtnValidation := bench.Operator.JoyBtnRaw);
ADVANCE_TIME(10000000);
bench(M1_PresetTriggerCmd := encoderM1.HwOut.PresetTriggerCmd, M1_PresetValueOut := encoderM1.HwOut.PresetValueOut, M2_PresetTriggerCmd := encoderM2.HwOut.PresetTriggerCmd, M2_PresetValueOut := encoderM2.HwOut.PresetValueOut, RawPosM1 := raw1, RawPosM2 := raw2); raw1 := bench.RawPosM1; raw2 := bench.RawPosM2;
hw1.RawPosIn := bench.Winch.COD1_PosValue; hw1.SlaveOperational := TRUE; hw2.RawPosIn := bench.Winch.COD2_PosValue; hw2.SlaveOperational := TRUE;
encoderM1(Enable := TRUE, HomingPermit := TRUE, HomingAtTargetM := btnM1, CfgHomingTargetM := 8.7, CfgTopSensorPosM := 8.7, HwIn := hw1, Cfg := cfgEncoder, Calib := calibM1); calibM1 := encoderM1.Calib;
bucketEdge(CLK := btnBucket);
encoderM2(Enable := TRUE, HomingPermit := TRUE, HomingAtTargetM := btnM2 OR bucketEdge.Q, CfgHomingTargetM := 23.7, CfgTopSensorPosM := 23.7, UseDynamicTarget := bucketEdge.Q, DynamicHomingTargetM := encoderM1.Measurement.CablePosM + cfgBucket.OffsetCloseM, HwIn := hw2, Cfg := cfgEncoder, Calib := calibM2); calibM2 := encoderM2.Calib;
bucket(Enable := TRUE, Mode := E_Mode.MAINT_N2, PowerContactorEngaged := TRUE, CablePosM1 := encoderM1.Measurement.CablePosM, CablePosM2 := encoderM2.Measurement.CablePosM, HomedM1 := encoderM1.Homed, HomedM2 := encoderM2.Homed, HomedAndReliableM1 := encoderM1.HomedAndReliable, HomedAndReliableM2 := encoderM2.HomedAndReliable, HomingSuspectM1 := encoderM1.HomingSuspect, HomingSuspectM2 := encoderM2.HomingSuspect, ConfirmClosePosition := btnBucket, Config := cfgBucket, BucketState := bucketState); bucketState := bucket.BucketState;
home.M1Status.HomedAndReliable := encoderM1.HomedAndReliable; home.M2Status.HomedAndReliable := encoderM2.HomedAndReliable; home(BucketOffsetValid := bucketState.BucketReferenced, BtnValidation := bench.Operator.JoyBtnRaw);
ADVANCE_TIME(10000000);
bench(M1_PresetTriggerCmd := encoderM1.HwOut.PresetTriggerCmd, M1_PresetValueOut := encoderM1.HwOut.PresetValueOut, M2_PresetTriggerCmd := encoderM2.HwOut.PresetTriggerCmd, M2_PresetValueOut := encoderM2.HwOut.PresetValueOut, RawPosM1 := raw1, RawPosM2 := raw2); raw1 := bench.RawPosM1; raw2 := bench.RawPosM2;
hw1.RawPosIn := bench.Winch.COD1_PosValue; hw1.SlaveOperational := TRUE; hw2.RawPosIn := bench.Winch.COD2_PosValue; hw2.SlaveOperational := TRUE;
encoderM1(Enable := TRUE, HomingPermit := TRUE, HomingAtTargetM := btnM1, CfgHomingTargetM := 8.7, CfgTopSensorPosM := 8.7, HwIn := hw1, Cfg := cfgEncoder, Calib := calibM1); calibM1 := encoderM1.Calib;
bucketEdge(CLK := btnBucket);
encoderM2(Enable := TRUE, HomingPermit := TRUE, HomingAtTargetM := btnM2 OR bucketEdge.Q, CfgHomingTargetM := 23.7, CfgTopSensorPosM := 23.7, UseDynamicTarget := bucketEdge.Q, DynamicHomingTargetM := encoderM1.Measurement.CablePosM + cfgBucket.OffsetCloseM, HwIn := hw2, Cfg := cfgEncoder, Calib := calibM2); calibM2 := encoderM2.Calib;
bucket(Enable := TRUE, Mode := E_Mode.MAINT_N2, PowerContactorEngaged := TRUE, CablePosM1 := encoderM1.Measurement.CablePosM, CablePosM2 := encoderM2.Measurement.CablePosM, HomedM1 := encoderM1.Homed, HomedM2 := encoderM2.Homed, HomedAndReliableM1 := encoderM1.HomedAndReliable, HomedAndReliableM2 := encoderM2.HomedAndReliable, HomingSuspectM1 := encoderM1.HomingSuspect, HomingSuspectM2 := encoderM2.HomingSuspect, ConfirmClosePosition := btnBucket, Config := cfgBucket, BucketState := bucketState); bucketState := bucket.BucketState;
home.M1Status.HomedAndReliable := encoderM1.HomedAndReliable; home.M2Status.HomedAndReliable := encoderM2.HomedAndReliable; home(BucketOffsetValid := bucketState.BucketReferenced, BtnValidation := bench.Operator.JoyBtnRaw);
ADVANCE_TIME(10000000);
bench(M1_PresetTriggerCmd := encoderM1.HwOut.PresetTriggerCmd, M1_PresetValueOut := encoderM1.HwOut.PresetValueOut, M2_PresetTriggerCmd := encoderM2.HwOut.PresetTriggerCmd, M2_PresetValueOut := encoderM2.HwOut.PresetValueOut, RawPosM1 := raw1, RawPosM2 := raw2); raw1 := bench.RawPosM1; raw2 := bench.RawPosM2;
hw1.RawPosIn := bench.Winch.COD1_PosValue; hw1.SlaveOperational := TRUE; hw2.RawPosIn := bench.Winch.COD2_PosValue; hw2.SlaveOperational := TRUE;
encoderM1(Enable := TRUE, HomingPermit := TRUE, HomingAtTargetM := btnM1, CfgHomingTargetM := 8.7, CfgTopSensorPosM := 8.7, HwIn := hw1, Cfg := cfgEncoder, Calib := calibM1); calibM1 := encoderM1.Calib;
bucketEdge(CLK := btnBucket);
encoderM2(Enable := TRUE, HomingPermit := TRUE, HomingAtTargetM := btnM2 OR bucketEdge.Q, CfgHomingTargetM := 23.7, CfgTopSensorPosM := 23.7, UseDynamicTarget := bucketEdge.Q, DynamicHomingTargetM := encoderM1.Measurement.CablePosM + cfgBucket.OffsetCloseM, HwIn := hw2, Cfg := cfgEncoder, Calib := calibM2); calibM2 := encoderM2.Calib;
bucket(Enable := TRUE, Mode := E_Mode.MAINT_N2, PowerContactorEngaged := TRUE, CablePosM1 := encoderM1.Measurement.CablePosM, CablePosM2 := encoderM2.Measurement.CablePosM, HomedM1 := encoderM1.Homed, HomedM2 := encoderM2.Homed, HomedAndReliableM1 := encoderM1.HomedAndReliable, HomedAndReliableM2 := encoderM2.HomedAndReliable, HomingSuspectM1 := encoderM1.HomingSuspect, HomingSuspectM2 := encoderM2.HomingSuspect, ConfirmClosePosition := btnBucket, Config := cfgBucket, BucketState := bucketState); bucketState := bucket.BucketState;
home.M1Status.HomedAndReliable := encoderM1.HomedAndReliable; home.M2Status.HomedAndReliable := encoderM2.HomedAndReliable; home(BucketOffsetValid := bucketState.BucketReferenced, BtnValidation := bench.Operator.JoyBtnRaw);
ADVANCE_TIME(10000000);
bench(M1_PresetTriggerCmd := encoderM1.HwOut.PresetTriggerCmd, M1_PresetValueOut := encoderM1.HwOut.PresetValueOut, M2_PresetTriggerCmd := encoderM2.HwOut.PresetTriggerCmd, M2_PresetValueOut := encoderM2.HwOut.PresetValueOut, RawPosM1 := raw1, RawPosM2 := raw2); raw1 := bench.RawPosM1; raw2 := bench.RawPosM2;
hw1.RawPosIn := bench.Winch.COD1_PosValue; hw1.SlaveOperational := TRUE; hw2.RawPosIn := bench.Winch.COD2_PosValue; hw2.SlaveOperational := TRUE;
encoderM1(Enable := TRUE, HomingPermit := TRUE, HomingAtTargetM := btnM1, CfgHomingTargetM := 8.7, CfgTopSensorPosM := 8.7, HwIn := hw1, Cfg := cfgEncoder, Calib := calibM1); calibM1 := encoderM1.Calib;
bucketEdge(CLK := btnBucket);
encoderM2(Enable := TRUE, HomingPermit := TRUE, HomingAtTargetM := btnM2 OR bucketEdge.Q, CfgHomingTargetM := 23.7, CfgTopSensorPosM := 23.7, UseDynamicTarget := bucketEdge.Q, DynamicHomingTargetM := encoderM1.Measurement.CablePosM + cfgBucket.OffsetCloseM, HwIn := hw2, Cfg := cfgEncoder, Calib := calibM2); calibM2 := encoderM2.Calib;
bucket(Enable := TRUE, Mode := E_Mode.MAINT_N2, PowerContactorEngaged := TRUE, CablePosM1 := encoderM1.Measurement.CablePosM, CablePosM2 := encoderM2.Measurement.CablePosM, HomedM1 := encoderM1.Homed, HomedM2 := encoderM2.Homed, HomedAndReliableM1 := encoderM1.HomedAndReliable, HomedAndReliableM2 := encoderM2.HomedAndReliable, HomingSuspectM1 := encoderM1.HomingSuspect, HomingSuspectM2 := encoderM2.HomingSuspect, ConfirmClosePosition := btnBucket, Config := cfgBucket, BucketState := bucketState); bucketState := bucket.BucketState;
home.M1Status.HomedAndReliable := encoderM1.HomedAndReliable; home.M2Status.HomedAndReliable := encoderM2.HomedAndReliable; home(BucketOffsetValid := bucketState.BucketReferenced, BtnValidation := bench.Operator.JoyBtnRaw);
ADVANCE_TIME(10000000);
bench(M1_PresetTriggerCmd := encoderM1.HwOut.PresetTriggerCmd, M1_PresetValueOut := encoderM1.HwOut.PresetValueOut, M2_PresetTriggerCmd := encoderM2.HwOut.PresetTriggerCmd, M2_PresetValueOut := encoderM2.HwOut.PresetValueOut, RawPosM1 := raw1, RawPosM2 := raw2); raw1 := bench.RawPosM1; raw2 := bench.RawPosM2;
hw1.RawPosIn := bench.Winch.COD1_PosValue; hw1.SlaveOperational := TRUE; hw2.RawPosIn := bench.Winch.COD2_PosValue; hw2.SlaveOperational := TRUE;
encoderM1(Enable := TRUE, HomingPermit := TRUE, HomingAtTargetM := btnM1, CfgHomingTargetM := 8.7, CfgTopSensorPosM := 8.7, HwIn := hw1, Cfg := cfgEncoder, Calib := calibM1); calibM1 := encoderM1.Calib;
bucketEdge(CLK := btnBucket);
encoderM2(Enable := TRUE, HomingPermit := TRUE, HomingAtTargetM := btnM2 OR bucketEdge.Q, CfgHomingTargetM := 23.7, CfgTopSensorPosM := 23.7, UseDynamicTarget := bucketEdge.Q, DynamicHomingTargetM := encoderM1.Measurement.CablePosM + cfgBucket.OffsetCloseM, HwIn := hw2, Cfg := cfgEncoder, Calib := calibM2); calibM2 := encoderM2.Calib;
bucket(Enable := TRUE, Mode := E_Mode.MAINT_N2, PowerContactorEngaged := TRUE, CablePosM1 := encoderM1.Measurement.CablePosM, CablePosM2 := encoderM2.Measurement.CablePosM, HomedM1 := encoderM1.Homed, HomedM2 := encoderM2.Homed, HomedAndReliableM1 := encoderM1.HomedAndReliable, HomedAndReliableM2 := encoderM2.HomedAndReliable, HomingSuspectM1 := encoderM1.HomingSuspect, HomingSuspectM2 := encoderM2.HomingSuspect, ConfirmClosePosition := btnBucket, Config := cfgBucket, BucketState := bucketState); bucketState := bucket.BucketState;
home.M1Status.HomedAndReliable := encoderM1.HomedAndReliable; home.M2Status.HomedAndReliable := encoderM2.HomedAndReliable; home(BucketOffsetValid := bucketState.BucketReferenced, BtnValidation := bench.Operator.JoyBtnRaw);
ADVANCE_TIME(10000000);
bench(M1_PresetTriggerCmd := encoderM1.HwOut.PresetTriggerCmd, M1_PresetValueOut := encoderM1.HwOut.PresetValueOut, M2_PresetTriggerCmd := encoderM2.HwOut.PresetTriggerCmd, M2_PresetValueOut := encoderM2.HwOut.PresetValueOut, RawPosM1 := raw1, RawPosM2 := raw2); raw1 := bench.RawPosM1; raw2 := bench.RawPosM2;
hw1.RawPosIn := bench.Winch.COD1_PosValue; hw1.SlaveOperational := TRUE; hw2.RawPosIn := bench.Winch.COD2_PosValue; hw2.SlaveOperational := TRUE;
encoderM1(Enable := TRUE, HomingPermit := TRUE, HomingAtTargetM := btnM1, CfgHomingTargetM := 8.7, CfgTopSensorPosM := 8.7, HwIn := hw1, Cfg := cfgEncoder, Calib := calibM1); calibM1 := encoderM1.Calib;
bucketEdge(CLK := btnBucket);
encoderM2(Enable := TRUE, HomingPermit := TRUE, HomingAtTargetM := btnM2 OR bucketEdge.Q, CfgHomingTargetM := 23.7, CfgTopSensorPosM := 23.7, UseDynamicTarget := bucketEdge.Q, DynamicHomingTargetM := encoderM1.Measurement.CablePosM + cfgBucket.OffsetCloseM, HwIn := hw2, Cfg := cfgEncoder, Calib := calibM2); calibM2 := encoderM2.Calib;
bucket(Enable := TRUE, Mode := E_Mode.MAINT_N2, PowerContactorEngaged := TRUE, CablePosM1 := encoderM1.Measurement.CablePosM, CablePosM2 := encoderM2.Measurement.CablePosM, HomedM1 := encoderM1.Homed, HomedM2 := encoderM2.Homed, HomedAndReliableM1 := encoderM1.HomedAndReliable, HomedAndReliableM2 := encoderM2.HomedAndReliable, HomingSuspectM1 := encoderM1.HomingSuspect, HomingSuspectM2 := encoderM2.HomingSuspect, ConfirmClosePosition := btnBucket, Config := cfgBucket, BucketState := bucketState); bucketState := bucket.BucketState;
home.M1Status.HomedAndReliable := encoderM1.HomedAndReliable; home.M2Status.HomedAndReliable := encoderM2.HomedAndReliable; home(BucketOffsetValid := bucketState.BucketReferenced, BtnValidation := bench.Operator.JoyBtnRaw);
ADVANCE_TIME(10000000);
bench(M1_PresetTriggerCmd := encoderM1.HwOut.PresetTriggerCmd, M1_PresetValueOut := encoderM1.HwOut.PresetValueOut, M2_PresetTriggerCmd := encoderM2.HwOut.PresetTriggerCmd, M2_PresetValueOut := encoderM2.HwOut.PresetValueOut, RawPosM1 := raw1, RawPosM2 := raw2); raw1 := bench.RawPosM1; raw2 := bench.RawPosM2;
hw1.RawPosIn := bench.Winch.COD1_PosValue; hw1.SlaveOperational := TRUE; hw2.RawPosIn := bench.Winch.COD2_PosValue; hw2.SlaveOperational := TRUE;
encoderM1(Enable := TRUE, HomingPermit := TRUE, HomingAtTargetM := btnM1, CfgHomingTargetM := 8.7, CfgTopSensorPosM := 8.7, HwIn := hw1, Cfg := cfgEncoder, Calib := calibM1); calibM1 := encoderM1.Calib;
bucketEdge(CLK := btnBucket);
encoderM2(Enable := TRUE, HomingPermit := TRUE, HomingAtTargetM := btnM2 OR bucketEdge.Q, CfgHomingTargetM := 23.7, CfgTopSensorPosM := 23.7, UseDynamicTarget := bucketEdge.Q, DynamicHomingTargetM := encoderM1.Measurement.CablePosM + cfgBucket.OffsetCloseM, HwIn := hw2, Cfg := cfgEncoder, Calib := calibM2); calibM2 := encoderM2.Calib;
bucket(Enable := TRUE, Mode := E_Mode.MAINT_N2, PowerContactorEngaged := TRUE, CablePosM1 := encoderM1.Measurement.CablePosM, CablePosM2 := encoderM2.Measurement.CablePosM, HomedM1 := encoderM1.Homed, HomedM2 := encoderM2.Homed, HomedAndReliableM1 := encoderM1.HomedAndReliable, HomedAndReliableM2 := encoderM2.HomedAndReliable, HomingSuspectM1 := encoderM1.HomingSuspect, HomingSuspectM2 := encoderM2.HomingSuspect, ConfirmClosePosition := btnBucket, Config := cfgBucket, BucketState := bucketState); bucketState := bucket.BucketState;
home.M1Status.HomedAndReliable := encoderM1.HomedAndReliable; home.M2Status.HomedAndReliable := encoderM2.HomedAndReliable; home(BucketOffsetValid := bucketState.BucketReferenced, BtnValidation := bench.Operator.JoyBtnRaw);
ADVANCE_TIME(10000000);
bench(M1_PresetTriggerCmd := encoderM1.HwOut.PresetTriggerCmd, M1_PresetValueOut := encoderM1.HwOut.PresetValueOut, M2_PresetTriggerCmd := encoderM2.HwOut.PresetTriggerCmd, M2_PresetValueOut := encoderM2.HwOut.PresetValueOut, RawPosM1 := raw1, RawPosM2 := raw2); raw1 := bench.RawPosM1; raw2 := bench.RawPosM2;
hw1.RawPosIn := bench.Winch.COD1_PosValue; hw1.SlaveOperational := TRUE; hw2.RawPosIn := bench.Winch.COD2_PosValue; hw2.SlaveOperational := TRUE;
encoderM1(Enable := TRUE, HomingPermit := TRUE, HomingAtTargetM := btnM1, CfgHomingTargetM := 8.7, CfgTopSensorPosM := 8.7, HwIn := hw1, Cfg := cfgEncoder, Calib := calibM1); calibM1 := encoderM1.Calib;
bucketEdge(CLK := btnBucket);
encoderM2(Enable := TRUE, HomingPermit := TRUE, HomingAtTargetM := btnM2 OR bucketEdge.Q, CfgHomingTargetM := 23.7, CfgTopSensorPosM := 23.7, UseDynamicTarget := bucketEdge.Q, DynamicHomingTargetM := encoderM1.Measurement.CablePosM + cfgBucket.OffsetCloseM, HwIn := hw2, Cfg := cfgEncoder, Calib := calibM2); calibM2 := encoderM2.Calib;
bucket(Enable := TRUE, Mode := E_Mode.MAINT_N2, PowerContactorEngaged := TRUE, CablePosM1 := encoderM1.Measurement.CablePosM, CablePosM2 := encoderM2.Measurement.CablePosM, HomedM1 := encoderM1.Homed, HomedM2 := encoderM2.Homed, HomedAndReliableM1 := encoderM1.HomedAndReliable, HomedAndReliableM2 := encoderM2.HomedAndReliable, HomingSuspectM1 := encoderM1.HomingSuspect, HomingSuspectM2 := encoderM2.HomingSuspect, ConfirmClosePosition := btnBucket, Config := cfgBucket, BucketState := bucketState); bucketState := bucket.BucketState;
home.M1Status.HomedAndReliable := encoderM1.HomedAndReliable; home.M2Status.HomedAndReliable := encoderM2.HomedAndReliable; home(BucketOffsetValid := bucketState.BucketReferenced, BtnValidation := bench.Operator.JoyBtnRaw);
ADVANCE_TIME(10000000);
bench(M1_PresetTriggerCmd := encoderM1.HwOut.PresetTriggerCmd, M1_PresetValueOut := encoderM1.HwOut.PresetValueOut, M2_PresetTriggerCmd := encoderM2.HwOut.PresetTriggerCmd, M2_PresetValueOut := encoderM2.HwOut.PresetValueOut, RawPosM1 := raw1, RawPosM2 := raw2); raw1 := bench.RawPosM1; raw2 := bench.RawPosM2;
hw1.RawPosIn := bench.Winch.COD1_PosValue; hw1.SlaveOperational := TRUE; hw2.RawPosIn := bench.Winch.COD2_PosValue; hw2.SlaveOperational := TRUE;
encoderM1(Enable := TRUE, HomingPermit := TRUE, HomingAtTargetM := btnM1, CfgHomingTargetM := 8.7, CfgTopSensorPosM := 8.7, HwIn := hw1, Cfg := cfgEncoder, Calib := calibM1); calibM1 := encoderM1.Calib;
bucketEdge(CLK := btnBucket);
encoderM2(Enable := TRUE, HomingPermit := TRUE, HomingAtTargetM := btnM2 OR bucketEdge.Q, CfgHomingTargetM := 23.7, CfgTopSensorPosM := 23.7, UseDynamicTarget := bucketEdge.Q, DynamicHomingTargetM := encoderM1.Measurement.CablePosM + cfgBucket.OffsetCloseM, HwIn := hw2, Cfg := cfgEncoder, Calib := calibM2); calibM2 := encoderM2.Calib;
bucket(Enable := TRUE, Mode := E_Mode.MAINT_N2, PowerContactorEngaged := TRUE, CablePosM1 := encoderM1.Measurement.CablePosM, CablePosM2 := encoderM2.Measurement.CablePosM, HomedM1 := encoderM1.Homed, HomedM2 := encoderM2.Homed, HomedAndReliableM1 := encoderM1.HomedAndReliable, HomedAndReliableM2 := encoderM2.HomedAndReliable, HomingSuspectM1 := encoderM1.HomingSuspect, HomingSuspectM2 := encoderM2.HomingSuspect, ConfirmClosePosition := btnBucket, Config := cfgBucket, BucketState := bucketState); bucketState := bucket.BucketState;
home.M1Status.HomedAndReliable := encoderM1.HomedAndReliable; home.M2Status.HomedAndReliable := encoderM2.HomedAndReliable; home(BucketOffsetValid := bucketState.BucketReferenced, BtnValidation := bench.Operator.JoyBtnRaw);
ADVANCE_TIME(10000000);
bench(M1_PresetTriggerCmd := encoderM1.HwOut.PresetTriggerCmd, M1_PresetValueOut := encoderM1.HwOut.PresetValueOut, M2_PresetTriggerCmd := encoderM2.HwOut.PresetTriggerCmd, M2_PresetValueOut := encoderM2.HwOut.PresetValueOut, RawPosM1 := raw1, RawPosM2 := raw2); raw1 := bench.RawPosM1; raw2 := bench.RawPosM2;
hw1.RawPosIn := bench.Winch.COD1_PosValue; hw1.SlaveOperational := TRUE; hw2.RawPosIn := bench.Winch.COD2_PosValue; hw2.SlaveOperational := TRUE;
encoderM1(Enable := TRUE, HomingPermit := TRUE, HomingAtTargetM := btnM1, CfgHomingTargetM := 8.7, CfgTopSensorPosM := 8.7, HwIn := hw1, Cfg := cfgEncoder, Calib := calibM1); calibM1 := encoderM1.Calib;
bucketEdge(CLK := btnBucket);
encoderM2(Enable := TRUE, HomingPermit := TRUE, HomingAtTargetM := btnM2 OR bucketEdge.Q, CfgHomingTargetM := 23.7, CfgTopSensorPosM := 23.7, UseDynamicTarget := bucketEdge.Q, DynamicHomingTargetM := encoderM1.Measurement.CablePosM + cfgBucket.OffsetCloseM, HwIn := hw2, Cfg := cfgEncoder, Calib := calibM2); calibM2 := encoderM2.Calib;
bucket(Enable := TRUE, Mode := E_Mode.MAINT_N2, PowerContactorEngaged := TRUE, CablePosM1 := encoderM1.Measurement.CablePosM, CablePosM2 := encoderM2.Measurement.CablePosM, HomedM1 := encoderM1.Homed, HomedM2 := encoderM2.Homed, HomedAndReliableM1 := encoderM1.HomedAndReliable, HomedAndReliableM2 := encoderM2.HomedAndReliable, HomingSuspectM1 := encoderM1.HomingSuspect, HomingSuspectM2 := encoderM2.HomingSuspect, ConfirmClosePosition := btnBucket, Config := cfgBucket, BucketState := bucketState); bucketState := bucket.BucketState;
home.M1Status.HomedAndReliable := encoderM1.HomedAndReliable; home.M2Status.HomedAndReliable := encoderM2.HomedAndReliable; home(BucketOffsetValid := bucketState.BucketReferenced, BtnValidation := bench.Operator.JoyBtnRaw);
ADVANCE_TIME(10000000);
bench(M1_PresetTriggerCmd := encoderM1.HwOut.PresetTriggerCmd, M1_PresetValueOut := encoderM1.HwOut.PresetValueOut, M2_PresetTriggerCmd := encoderM2.HwOut.PresetTriggerCmd, M2_PresetValueOut := encoderM2.HwOut.PresetValueOut, RawPosM1 := raw1, RawPosM2 := raw2); raw1 := bench.RawPosM1; raw2 := bench.RawPosM2;
hw1.RawPosIn := bench.Winch.COD1_PosValue; hw1.SlaveOperational := TRUE; hw2.RawPosIn := bench.Winch.COD2_PosValue; hw2.SlaveOperational := TRUE;
encoderM1(Enable := TRUE, HomingPermit := TRUE, HomingAtTargetM := btnM1, CfgHomingTargetM := 8.7, CfgTopSensorPosM := 8.7, HwIn := hw1, Cfg := cfgEncoder, Calib := calibM1); calibM1 := encoderM1.Calib;
bucketEdge(CLK := btnBucket);
encoderM2(Enable := TRUE, HomingPermit := TRUE, HomingAtTargetM := btnM2 OR bucketEdge.Q, CfgHomingTargetM := 23.7, CfgTopSensorPosM := 23.7, UseDynamicTarget := bucketEdge.Q, DynamicHomingTargetM := encoderM1.Measurement.CablePosM + cfgBucket.OffsetCloseM, HwIn := hw2, Cfg := cfgEncoder, Calib := calibM2); calibM2 := encoderM2.Calib;
bucket(Enable := TRUE, Mode := E_Mode.MAINT_N2, PowerContactorEngaged := TRUE, CablePosM1 := encoderM1.Measurement.CablePosM, CablePosM2 := encoderM2.Measurement.CablePosM, HomedM1 := encoderM1.Homed, HomedM2 := encoderM2.Homed, HomedAndReliableM1 := encoderM1.HomedAndReliable, HomedAndReliableM2 := encoderM2.HomedAndReliable, HomingSuspectM1 := encoderM1.HomingSuspect, HomingSuspectM2 := encoderM2.HomingSuspect, ConfirmClosePosition := btnBucket, Config := cfgBucket, BucketState := bucketState); bucketState := bucket.BucketState;
home.M1Status.HomedAndReliable := encoderM1.HomedAndReliable; home.M2Status.HomedAndReliable := encoderM2.HomedAndReliable; home(BucketOffsetValid := bucketState.BucketReferenced, BtnValidation := bench.Operator.JoyBtnRaw);
ADVANCE_TIME(10000000);
bench(M1_PresetTriggerCmd := encoderM1.HwOut.PresetTriggerCmd, M1_PresetValueOut := encoderM1.HwOut.PresetValueOut, M2_PresetTriggerCmd := encoderM2.HwOut.PresetTriggerCmd, M2_PresetValueOut := encoderM2.HwOut.PresetValueOut, RawPosM1 := raw1, RawPosM2 := raw2); raw1 := bench.RawPosM1; raw2 := bench.RawPosM2;
hw1.RawPosIn := bench.Winch.COD1_PosValue; hw1.SlaveOperational := TRUE; hw2.RawPosIn := bench.Winch.COD2_PosValue; hw2.SlaveOperational := TRUE;
encoderM1(Enable := TRUE, HomingPermit := TRUE, HomingAtTargetM := btnM1, CfgHomingTargetM := 8.7, CfgTopSensorPosM := 8.7, HwIn := hw1, Cfg := cfgEncoder, Calib := calibM1); calibM1 := encoderM1.Calib;
bucketEdge(CLK := btnBucket);
encoderM2(Enable := TRUE, HomingPermit := TRUE, HomingAtTargetM := btnM2 OR bucketEdge.Q, CfgHomingTargetM := 23.7, CfgTopSensorPosM := 23.7, UseDynamicTarget := bucketEdge.Q, DynamicHomingTargetM := encoderM1.Measurement.CablePosM + cfgBucket.OffsetCloseM, HwIn := hw2, Cfg := cfgEncoder, Calib := calibM2); calibM2 := encoderM2.Calib;
bucket(Enable := TRUE, Mode := E_Mode.MAINT_N2, PowerContactorEngaged := TRUE, CablePosM1 := encoderM1.Measurement.CablePosM, CablePosM2 := encoderM2.Measurement.CablePosM, HomedM1 := encoderM1.Homed, HomedM2 := encoderM2.Homed, HomedAndReliableM1 := encoderM1.HomedAndReliable, HomedAndReliableM2 := encoderM2.HomedAndReliable, HomingSuspectM1 := encoderM1.HomingSuspect, HomingSuspectM2 := encoderM2.HomingSuspect, ConfirmClosePosition := btnBucket, Config := cfgBucket, BucketState := bucketState); bucketState := bucket.BucketState;
home.M1Status.HomedAndReliable := encoderM1.HomedAndReliable; home.M2Status.HomedAndReliable := encoderM2.HomedAndReliable; home(BucketOffsetValid := bucketState.BucketReferenced, BtnValidation := bench.Operator.JoyBtnRaw);
ADVANCE_TIME(10000000);
bench(M1_PresetTriggerCmd := encoderM1.HwOut.PresetTriggerCmd, M1_PresetValueOut := encoderM1.HwOut.PresetValueOut, M2_PresetTriggerCmd := encoderM2.HwOut.PresetTriggerCmd, M2_PresetValueOut := encoderM2.HwOut.PresetValueOut, RawPosM1 := raw1, RawPosM2 := raw2); raw1 := bench.RawPosM1; raw2 := bench.RawPosM2;
hw1.RawPosIn := bench.Winch.COD1_PosValue; hw1.SlaveOperational := TRUE; hw2.RawPosIn := bench.Winch.COD2_PosValue; hw2.SlaveOperational := TRUE;
encoderM1(Enable := TRUE, HomingPermit := TRUE, HomingAtTargetM := btnM1, CfgHomingTargetM := 8.7, CfgTopSensorPosM := 8.7, HwIn := hw1, Cfg := cfgEncoder, Calib := calibM1); calibM1 := encoderM1.Calib;
bucketEdge(CLK := btnBucket);
encoderM2(Enable := TRUE, HomingPermit := TRUE, HomingAtTargetM := btnM2 OR bucketEdge.Q, CfgHomingTargetM := 23.7, CfgTopSensorPosM := 23.7, UseDynamicTarget := bucketEdge.Q, DynamicHomingTargetM := encoderM1.Measurement.CablePosM + cfgBucket.OffsetCloseM, HwIn := hw2, Cfg := cfgEncoder, Calib := calibM2); calibM2 := encoderM2.Calib;
bucket(Enable := TRUE, Mode := E_Mode.MAINT_N2, PowerContactorEngaged := TRUE, CablePosM1 := encoderM1.Measurement.CablePosM, CablePosM2 := encoderM2.Measurement.CablePosM, HomedM1 := encoderM1.Homed, HomedM2 := encoderM2.Homed, HomedAndReliableM1 := encoderM1.HomedAndReliable, HomedAndReliableM2 := encoderM2.HomedAndReliable, HomingSuspectM1 := encoderM1.HomingSuspect, HomingSuspectM2 := encoderM2.HomingSuspect, ConfirmClosePosition := btnBucket, Config := cfgBucket, BucketState := bucketState); bucketState := bucket.BucketState;
home.M1Status.HomedAndReliable := encoderM1.HomedAndReliable; home.M2Status.HomedAndReliable := encoderM2.HomedAndReliable; home(BucketOffsetValid := bucketState.BucketReferenced, BtnValidation := bench.Operator.JoyBtnRaw);
ADVANCE_TIME(10000000);
bench(M1_PresetTriggerCmd := encoderM1.HwOut.PresetTriggerCmd, M1_PresetValueOut := encoderM1.HwOut.PresetValueOut, M2_PresetTriggerCmd := encoderM2.HwOut.PresetTriggerCmd, M2_PresetValueOut := encoderM2.HwOut.PresetValueOut, RawPosM1 := raw1, RawPosM2 := raw2); raw1 := bench.RawPosM1; raw2 := bench.RawPosM2;
hw1.RawPosIn := bench.Winch.COD1_PosValue; hw1.SlaveOperational := TRUE; hw2.RawPosIn := bench.Winch.COD2_PosValue; hw2.SlaveOperational := TRUE;
encoderM1(Enable := TRUE, HomingPermit := TRUE, HomingAtTargetM := btnM1, CfgHomingTargetM := 8.7, CfgTopSensorPosM := 8.7, HwIn := hw1, Cfg := cfgEncoder, Calib := calibM1); calibM1 := encoderM1.Calib;
bucketEdge(CLK := btnBucket);
encoderM2(Enable := TRUE, HomingPermit := TRUE, HomingAtTargetM := btnM2 OR bucketEdge.Q, CfgHomingTargetM := 23.7, CfgTopSensorPosM := 23.7, UseDynamicTarget := bucketEdge.Q, DynamicHomingTargetM := encoderM1.Measurement.CablePosM + cfgBucket.OffsetCloseM, HwIn := hw2, Cfg := cfgEncoder, Calib := calibM2); calibM2 := encoderM2.Calib;
bucket(Enable := TRUE, Mode := E_Mode.MAINT_N2, PowerContactorEngaged := TRUE, CablePosM1 := encoderM1.Measurement.CablePosM, CablePosM2 := encoderM2.Measurement.CablePosM, HomedM1 := encoderM1.Homed, HomedM2 := encoderM2.Homed, HomedAndReliableM1 := encoderM1.HomedAndReliable, HomedAndReliableM2 := encoderM2.HomedAndReliable, HomingSuspectM1 := encoderM1.HomingSuspect, HomingSuspectM2 := encoderM2.HomingSuspect, ConfirmClosePosition := btnBucket, Config := cfgBucket, BucketState := bucketState); bucketState := bucket.BucketState;
home.M1Status.HomedAndReliable := encoderM1.HomedAndReliable; home.M2Status.HomedAndReliable := encoderM2.HomedAndReliable; home(BucketOffsetValid := bucketState.BucketReferenced, BtnValidation := bench.Operator.JoyBtnRaw);
ASSERT_TRUE(encoderM2.HomedAndReliable, 'Deuxieme bouton reference M2'); ASSERT_FALSE(home.MachineHomed, 'Machine attend reference benne');
btnBucket := TRUE;
ADVANCE_TIME(10000000);
bench(M1_PresetTriggerCmd := encoderM1.HwOut.PresetTriggerCmd, M1_PresetValueOut := encoderM1.HwOut.PresetValueOut, M2_PresetTriggerCmd := encoderM2.HwOut.PresetTriggerCmd, M2_PresetValueOut := encoderM2.HwOut.PresetValueOut, RawPosM1 := raw1, RawPosM2 := raw2); raw1 := bench.RawPosM1; raw2 := bench.RawPosM2;
hw1.RawPosIn := bench.Winch.COD1_PosValue; hw1.SlaveOperational := TRUE; hw2.RawPosIn := bench.Winch.COD2_PosValue; hw2.SlaveOperational := TRUE;
encoderM1(Enable := TRUE, HomingPermit := TRUE, HomingAtTargetM := btnM1, CfgHomingTargetM := 8.7, CfgTopSensorPosM := 8.7, HwIn := hw1, Cfg := cfgEncoder, Calib := calibM1); calibM1 := encoderM1.Calib;
bucketEdge(CLK := btnBucket);
encoderM2(Enable := TRUE, HomingPermit := TRUE, HomingAtTargetM := btnM2 OR bucketEdge.Q, CfgHomingTargetM := 23.7, CfgTopSensorPosM := 23.7, UseDynamicTarget := bucketEdge.Q, DynamicHomingTargetM := encoderM1.Measurement.CablePosM + cfgBucket.OffsetCloseM, HwIn := hw2, Cfg := cfgEncoder, Calib := calibM2); calibM2 := encoderM2.Calib;
bucket(Enable := TRUE, Mode := E_Mode.MAINT_N2, PowerContactorEngaged := TRUE, CablePosM1 := encoderM1.Measurement.CablePosM, CablePosM2 := encoderM2.Measurement.CablePosM, HomedM1 := encoderM1.Homed, HomedM2 := encoderM2.Homed, HomedAndReliableM1 := encoderM1.HomedAndReliable, HomedAndReliableM2 := encoderM2.HomedAndReliable, HomingSuspectM1 := encoderM1.HomingSuspect, HomingSuspectM2 := encoderM2.HomingSuspect, ConfirmClosePosition := btnBucket, Config := cfgBucket, BucketState := bucketState); bucketState := bucket.BucketState;
home.M1Status.HomedAndReliable := encoderM1.HomedAndReliable; home.M2Status.HomedAndReliable := encoderM2.HomedAndReliable; home(BucketOffsetValid := bucketState.BucketReferenced, BtnValidation := bench.Operator.JoyBtnRaw);
btnBucket := FALSE;
ADVANCE_TIME(10000000);
bench(M1_PresetTriggerCmd := encoderM1.HwOut.PresetTriggerCmd, M1_PresetValueOut := encoderM1.HwOut.PresetValueOut, M2_PresetTriggerCmd := encoderM2.HwOut.PresetTriggerCmd, M2_PresetValueOut := encoderM2.HwOut.PresetValueOut, RawPosM1 := raw1, RawPosM2 := raw2); raw1 := bench.RawPosM1; raw2 := bench.RawPosM2;
hw1.RawPosIn := bench.Winch.COD1_PosValue; hw1.SlaveOperational := TRUE; hw2.RawPosIn := bench.Winch.COD2_PosValue; hw2.SlaveOperational := TRUE;
encoderM1(Enable := TRUE, HomingPermit := TRUE, HomingAtTargetM := btnM1, CfgHomingTargetM := 8.7, CfgTopSensorPosM := 8.7, HwIn := hw1, Cfg := cfgEncoder, Calib := calibM1); calibM1 := encoderM1.Calib;
bucketEdge(CLK := btnBucket);
encoderM2(Enable := TRUE, HomingPermit := TRUE, HomingAtTargetM := btnM2 OR bucketEdge.Q, CfgHomingTargetM := 23.7, CfgTopSensorPosM := 23.7, UseDynamicTarget := bucketEdge.Q, DynamicHomingTargetM := encoderM1.Measurement.CablePosM + cfgBucket.OffsetCloseM, HwIn := hw2, Cfg := cfgEncoder, Calib := calibM2); calibM2 := encoderM2.Calib;
bucket(Enable := TRUE, Mode := E_Mode.MAINT_N2, PowerContactorEngaged := TRUE, CablePosM1 := encoderM1.Measurement.CablePosM, CablePosM2 := encoderM2.Measurement.CablePosM, HomedM1 := encoderM1.Homed, HomedM2 := encoderM2.Homed, HomedAndReliableM1 := encoderM1.HomedAndReliable, HomedAndReliableM2 := encoderM2.HomedAndReliable, HomingSuspectM1 := encoderM1.HomingSuspect, HomingSuspectM2 := encoderM2.HomingSuspect, ConfirmClosePosition := btnBucket, Config := cfgBucket, BucketState := bucketState); bucketState := bucket.BucketState;
home.M1Status.HomedAndReliable := encoderM1.HomedAndReliable; home.M2Status.HomedAndReliable := encoderM2.HomedAndReliable; home(BucketOffsetValid := bucketState.BucketReferenced, BtnValidation := bench.Operator.JoyBtnRaw);
ADVANCE_TIME(10000000);
bench(M1_PresetTriggerCmd := encoderM1.HwOut.PresetTriggerCmd, M1_PresetValueOut := encoderM1.HwOut.PresetValueOut, M2_PresetTriggerCmd := encoderM2.HwOut.PresetTriggerCmd, M2_PresetValueOut := encoderM2.HwOut.PresetValueOut, RawPosM1 := raw1, RawPosM2 := raw2); raw1 := bench.RawPosM1; raw2 := bench.RawPosM2;
hw1.RawPosIn := bench.Winch.COD1_PosValue; hw1.SlaveOperational := TRUE; hw2.RawPosIn := bench.Winch.COD2_PosValue; hw2.SlaveOperational := TRUE;
encoderM1(Enable := TRUE, HomingPermit := TRUE, HomingAtTargetM := btnM1, CfgHomingTargetM := 8.7, CfgTopSensorPosM := 8.7, HwIn := hw1, Cfg := cfgEncoder, Calib := calibM1); calibM1 := encoderM1.Calib;
bucketEdge(CLK := btnBucket);
encoderM2(Enable := TRUE, HomingPermit := TRUE, HomingAtTargetM := btnM2 OR bucketEdge.Q, CfgHomingTargetM := 23.7, CfgTopSensorPosM := 23.7, UseDynamicTarget := bucketEdge.Q, DynamicHomingTargetM := encoderM1.Measurement.CablePosM + cfgBucket.OffsetCloseM, HwIn := hw2, Cfg := cfgEncoder, Calib := calibM2); calibM2 := encoderM2.Calib;
bucket(Enable := TRUE, Mode := E_Mode.MAINT_N2, PowerContactorEngaged := TRUE, CablePosM1 := encoderM1.Measurement.CablePosM, CablePosM2 := encoderM2.Measurement.CablePosM, HomedM1 := encoderM1.Homed, HomedM2 := encoderM2.Homed, HomedAndReliableM1 := encoderM1.HomedAndReliable, HomedAndReliableM2 := encoderM2.HomedAndReliable, HomingSuspectM1 := encoderM1.HomingSuspect, HomingSuspectM2 := encoderM2.HomingSuspect, ConfirmClosePosition := btnBucket, Config := cfgBucket, BucketState := bucketState); bucketState := bucket.BucketState;
home.M1Status.HomedAndReliable := encoderM1.HomedAndReliable; home.M2Status.HomedAndReliable := encoderM2.HomedAndReliable; home(BucketOffsetValid := bucketState.BucketReferenced, BtnValidation := bench.Operator.JoyBtnRaw);
ADVANCE_TIME(10000000);
bench(M1_PresetTriggerCmd := encoderM1.HwOut.PresetTriggerCmd, M1_PresetValueOut := encoderM1.HwOut.PresetValueOut, M2_PresetTriggerCmd := encoderM2.HwOut.PresetTriggerCmd, M2_PresetValueOut := encoderM2.HwOut.PresetValueOut, RawPosM1 := raw1, RawPosM2 := raw2); raw1 := bench.RawPosM1; raw2 := bench.RawPosM2;
hw1.RawPosIn := bench.Winch.COD1_PosValue; hw1.SlaveOperational := TRUE; hw2.RawPosIn := bench.Winch.COD2_PosValue; hw2.SlaveOperational := TRUE;
encoderM1(Enable := TRUE, HomingPermit := TRUE, HomingAtTargetM := btnM1, CfgHomingTargetM := 8.7, CfgTopSensorPosM := 8.7, HwIn := hw1, Cfg := cfgEncoder, Calib := calibM1); calibM1 := encoderM1.Calib;
bucketEdge(CLK := btnBucket);
encoderM2(Enable := TRUE, HomingPermit := TRUE, HomingAtTargetM := btnM2 OR bucketEdge.Q, CfgHomingTargetM := 23.7, CfgTopSensorPosM := 23.7, UseDynamicTarget := bucketEdge.Q, DynamicHomingTargetM := encoderM1.Measurement.CablePosM + cfgBucket.OffsetCloseM, HwIn := hw2, Cfg := cfgEncoder, Calib := calibM2); calibM2 := encoderM2.Calib;
bucket(Enable := TRUE, Mode := E_Mode.MAINT_N2, PowerContactorEngaged := TRUE, CablePosM1 := encoderM1.Measurement.CablePosM, CablePosM2 := encoderM2.Measurement.CablePosM, HomedM1 := encoderM1.Homed, HomedM2 := encoderM2.Homed, HomedAndReliableM1 := encoderM1.HomedAndReliable, HomedAndReliableM2 := encoderM2.HomedAndReliable, HomingSuspectM1 := encoderM1.HomingSuspect, HomingSuspectM2 := encoderM2.HomingSuspect, ConfirmClosePosition := btnBucket, Config := cfgBucket, BucketState := bucketState); bucketState := bucket.BucketState;
home.M1Status.HomedAndReliable := encoderM1.HomedAndReliable; home.M2Status.HomedAndReliable := encoderM2.HomedAndReliable; home(BucketOffsetValid := bucketState.BucketReferenced, BtnValidation := bench.Operator.JoyBtnRaw);
ADVANCE_TIME(10000000);
bench(M1_PresetTriggerCmd := encoderM1.HwOut.PresetTriggerCmd, M1_PresetValueOut := encoderM1.HwOut.PresetValueOut, M2_PresetTriggerCmd := encoderM2.HwOut.PresetTriggerCmd, M2_PresetValueOut := encoderM2.HwOut.PresetValueOut, RawPosM1 := raw1, RawPosM2 := raw2); raw1 := bench.RawPosM1; raw2 := bench.RawPosM2;
hw1.RawPosIn := bench.Winch.COD1_PosValue; hw1.SlaveOperational := TRUE; hw2.RawPosIn := bench.Winch.COD2_PosValue; hw2.SlaveOperational := TRUE;
encoderM1(Enable := TRUE, HomingPermit := TRUE, HomingAtTargetM := btnM1, CfgHomingTargetM := 8.7, CfgTopSensorPosM := 8.7, HwIn := hw1, Cfg := cfgEncoder, Calib := calibM1); calibM1 := encoderM1.Calib;
bucketEdge(CLK := btnBucket);
encoderM2(Enable := TRUE, HomingPermit := TRUE, HomingAtTargetM := btnM2 OR bucketEdge.Q, CfgHomingTargetM := 23.7, CfgTopSensorPosM := 23.7, UseDynamicTarget := bucketEdge.Q, DynamicHomingTargetM := encoderM1.Measurement.CablePosM + cfgBucket.OffsetCloseM, HwIn := hw2, Cfg := cfgEncoder, Calib := calibM2); calibM2 := encoderM2.Calib;
bucket(Enable := TRUE, Mode := E_Mode.MAINT_N2, PowerContactorEngaged := TRUE, CablePosM1 := encoderM1.Measurement.CablePosM, CablePosM2 := encoderM2.Measurement.CablePosM, HomedM1 := encoderM1.Homed, HomedM2 := encoderM2.Homed, HomedAndReliableM1 := encoderM1.HomedAndReliable, HomedAndReliableM2 := encoderM2.HomedAndReliable, HomingSuspectM1 := encoderM1.HomingSuspect, HomingSuspectM2 := encoderM2.HomingSuspect, ConfirmClosePosition := btnBucket, Config := cfgBucket, BucketState := bucketState); bucketState := bucket.BucketState;
home.M1Status.HomedAndReliable := encoderM1.HomedAndReliable; home.M2Status.HomedAndReliable := encoderM2.HomedAndReliable; home(BucketOffsetValid := bucketState.BucketReferenced, BtnValidation := bench.Operator.JoyBtnRaw);
ADVANCE_TIME(10000000);
bench(M1_PresetTriggerCmd := encoderM1.HwOut.PresetTriggerCmd, M1_PresetValueOut := encoderM1.HwOut.PresetValueOut, M2_PresetTriggerCmd := encoderM2.HwOut.PresetTriggerCmd, M2_PresetValueOut := encoderM2.HwOut.PresetValueOut, RawPosM1 := raw1, RawPosM2 := raw2); raw1 := bench.RawPosM1; raw2 := bench.RawPosM2;
hw1.RawPosIn := bench.Winch.COD1_PosValue; hw1.SlaveOperational := TRUE; hw2.RawPosIn := bench.Winch.COD2_PosValue; hw2.SlaveOperational := TRUE;
encoderM1(Enable := TRUE, HomingPermit := TRUE, HomingAtTargetM := btnM1, CfgHomingTargetM := 8.7, CfgTopSensorPosM := 8.7, HwIn := hw1, Cfg := cfgEncoder, Calib := calibM1); calibM1 := encoderM1.Calib;
bucketEdge(CLK := btnBucket);
encoderM2(Enable := TRUE, HomingPermit := TRUE, HomingAtTargetM := btnM2 OR bucketEdge.Q, CfgHomingTargetM := 23.7, CfgTopSensorPosM := 23.7, UseDynamicTarget := bucketEdge.Q, DynamicHomingTargetM := encoderM1.Measurement.CablePosM + cfgBucket.OffsetCloseM, HwIn := hw2, Cfg := cfgEncoder, Calib := calibM2); calibM2 := encoderM2.Calib;
bucket(Enable := TRUE, Mode := E_Mode.MAINT_N2, PowerContactorEngaged := TRUE, CablePosM1 := encoderM1.Measurement.CablePosM, CablePosM2 := encoderM2.Measurement.CablePosM, HomedM1 := encoderM1.Homed, HomedM2 := encoderM2.Homed, HomedAndReliableM1 := encoderM1.HomedAndReliable, HomedAndReliableM2 := encoderM2.HomedAndReliable, HomingSuspectM1 := encoderM1.HomingSuspect, HomingSuspectM2 := encoderM2.HomingSuspect, ConfirmClosePosition := btnBucket, Config := cfgBucket, BucketState := bucketState); bucketState := bucket.BucketState;
home.M1Status.HomedAndReliable := encoderM1.HomedAndReliable; home.M2Status.HomedAndReliable := encoderM2.HomedAndReliable; home(BucketOffsetValid := bucketState.BucketReferenced, BtnValidation := bench.Operator.JoyBtnRaw);
ADVANCE_TIME(10000000);
bench(M1_PresetTriggerCmd := encoderM1.HwOut.PresetTriggerCmd, M1_PresetValueOut := encoderM1.HwOut.PresetValueOut, M2_PresetTriggerCmd := encoderM2.HwOut.PresetTriggerCmd, M2_PresetValueOut := encoderM2.HwOut.PresetValueOut, RawPosM1 := raw1, RawPosM2 := raw2); raw1 := bench.RawPosM1; raw2 := bench.RawPosM2;
hw1.RawPosIn := bench.Winch.COD1_PosValue; hw1.SlaveOperational := TRUE; hw2.RawPosIn := bench.Winch.COD2_PosValue; hw2.SlaveOperational := TRUE;
encoderM1(Enable := TRUE, HomingPermit := TRUE, HomingAtTargetM := btnM1, CfgHomingTargetM := 8.7, CfgTopSensorPosM := 8.7, HwIn := hw1, Cfg := cfgEncoder, Calib := calibM1); calibM1 := encoderM1.Calib;
bucketEdge(CLK := btnBucket);
encoderM2(Enable := TRUE, HomingPermit := TRUE, HomingAtTargetM := btnM2 OR bucketEdge.Q, CfgHomingTargetM := 23.7, CfgTopSensorPosM := 23.7, UseDynamicTarget := bucketEdge.Q, DynamicHomingTargetM := encoderM1.Measurement.CablePosM + cfgBucket.OffsetCloseM, HwIn := hw2, Cfg := cfgEncoder, Calib := calibM2); calibM2 := encoderM2.Calib;
bucket(Enable := TRUE, Mode := E_Mode.MAINT_N2, PowerContactorEngaged := TRUE, CablePosM1 := encoderM1.Measurement.CablePosM, CablePosM2 := encoderM2.Measurement.CablePosM, HomedM1 := encoderM1.Homed, HomedM2 := encoderM2.Homed, HomedAndReliableM1 := encoderM1.HomedAndReliable, HomedAndReliableM2 := encoderM2.HomedAndReliable, HomingSuspectM1 := encoderM1.HomingSuspect, HomingSuspectM2 := encoderM2.HomingSuspect, ConfirmClosePosition := btnBucket, Config := cfgBucket, BucketState := bucketState); bucketState := bucket.BucketState;
home.M1Status.HomedAndReliable := encoderM1.HomedAndReliable; home.M2Status.HomedAndReliable := encoderM2.HomedAndReliable; home(BucketOffsetValid := bucketState.BucketReferenced, BtnValidation := bench.Operator.JoyBtnRaw);
ADVANCE_TIME(10000000);
bench(M1_PresetTriggerCmd := encoderM1.HwOut.PresetTriggerCmd, M1_PresetValueOut := encoderM1.HwOut.PresetValueOut, M2_PresetTriggerCmd := encoderM2.HwOut.PresetTriggerCmd, M2_PresetValueOut := encoderM2.HwOut.PresetValueOut, RawPosM1 := raw1, RawPosM2 := raw2); raw1 := bench.RawPosM1; raw2 := bench.RawPosM2;
hw1.RawPosIn := bench.Winch.COD1_PosValue; hw1.SlaveOperational := TRUE; hw2.RawPosIn := bench.Winch.COD2_PosValue; hw2.SlaveOperational := TRUE;
encoderM1(Enable := TRUE, HomingPermit := TRUE, HomingAtTargetM := btnM1, CfgHomingTargetM := 8.7, CfgTopSensorPosM := 8.7, HwIn := hw1, Cfg := cfgEncoder, Calib := calibM1); calibM1 := encoderM1.Calib;
bucketEdge(CLK := btnBucket);
encoderM2(Enable := TRUE, HomingPermit := TRUE, HomingAtTargetM := btnM2 OR bucketEdge.Q, CfgHomingTargetM := 23.7, CfgTopSensorPosM := 23.7, UseDynamicTarget := bucketEdge.Q, DynamicHomingTargetM := encoderM1.Measurement.CablePosM + cfgBucket.OffsetCloseM, HwIn := hw2, Cfg := cfgEncoder, Calib := calibM2); calibM2 := encoderM2.Calib;
bucket(Enable := TRUE, Mode := E_Mode.MAINT_N2, PowerContactorEngaged := TRUE, CablePosM1 := encoderM1.Measurement.CablePosM, CablePosM2 := encoderM2.Measurement.CablePosM, HomedM1 := encoderM1.Homed, HomedM2 := encoderM2.Homed, HomedAndReliableM1 := encoderM1.HomedAndReliable, HomedAndReliableM2 := encoderM2.HomedAndReliable, HomingSuspectM1 := encoderM1.HomingSuspect, HomingSuspectM2 := encoderM2.HomingSuspect, ConfirmClosePosition := btnBucket, Config := cfgBucket, BucketState := bucketState); bucketState := bucket.BucketState;
home.M1Status.HomedAndReliable := encoderM1.HomedAndReliable; home.M2Status.HomedAndReliable := encoderM2.HomedAndReliable; home(BucketOffsetValid := bucketState.BucketReferenced, BtnValidation := bench.Operator.JoyBtnRaw);
ADVANCE_TIME(10000000);
bench(M1_PresetTriggerCmd := encoderM1.HwOut.PresetTriggerCmd, M1_PresetValueOut := encoderM1.HwOut.PresetValueOut, M2_PresetTriggerCmd := encoderM2.HwOut.PresetTriggerCmd, M2_PresetValueOut := encoderM2.HwOut.PresetValueOut, RawPosM1 := raw1, RawPosM2 := raw2); raw1 := bench.RawPosM1; raw2 := bench.RawPosM2;
hw1.RawPosIn := bench.Winch.COD1_PosValue; hw1.SlaveOperational := TRUE; hw2.RawPosIn := bench.Winch.COD2_PosValue; hw2.SlaveOperational := TRUE;
encoderM1(Enable := TRUE, HomingPermit := TRUE, HomingAtTargetM := btnM1, CfgHomingTargetM := 8.7, CfgTopSensorPosM := 8.7, HwIn := hw1, Cfg := cfgEncoder, Calib := calibM1); calibM1 := encoderM1.Calib;
bucketEdge(CLK := btnBucket);
encoderM2(Enable := TRUE, HomingPermit := TRUE, HomingAtTargetM := btnM2 OR bucketEdge.Q, CfgHomingTargetM := 23.7, CfgTopSensorPosM := 23.7, UseDynamicTarget := bucketEdge.Q, DynamicHomingTargetM := encoderM1.Measurement.CablePosM + cfgBucket.OffsetCloseM, HwIn := hw2, Cfg := cfgEncoder, Calib := calibM2); calibM2 := encoderM2.Calib;
bucket(Enable := TRUE, Mode := E_Mode.MAINT_N2, PowerContactorEngaged := TRUE, CablePosM1 := encoderM1.Measurement.CablePosM, CablePosM2 := encoderM2.Measurement.CablePosM, HomedM1 := encoderM1.Homed, HomedM2 := encoderM2.Homed, HomedAndReliableM1 := encoderM1.HomedAndReliable, HomedAndReliableM2 := encoderM2.HomedAndReliable, HomingSuspectM1 := encoderM1.HomingSuspect, HomingSuspectM2 := encoderM2.HomingSuspect, ConfirmClosePosition := btnBucket, Config := cfgBucket, BucketState := bucketState); bucketState := bucket.BucketState;
home.M1Status.HomedAndReliable := encoderM1.HomedAndReliable; home.M2Status.HomedAndReliable := encoderM2.HomedAndReliable; home(BucketOffsetValid := bucketState.BucketReferenced, BtnValidation := bench.Operator.JoyBtnRaw);
ADVANCE_TIME(10000000);
bench(M1_PresetTriggerCmd := encoderM1.HwOut.PresetTriggerCmd, M1_PresetValueOut := encoderM1.HwOut.PresetValueOut, M2_PresetTriggerCmd := encoderM2.HwOut.PresetTriggerCmd, M2_PresetValueOut := encoderM2.HwOut.PresetValueOut, RawPosM1 := raw1, RawPosM2 := raw2); raw1 := bench.RawPosM1; raw2 := bench.RawPosM2;
hw1.RawPosIn := bench.Winch.COD1_PosValue; hw1.SlaveOperational := TRUE; hw2.RawPosIn := bench.Winch.COD2_PosValue; hw2.SlaveOperational := TRUE;
encoderM1(Enable := TRUE, HomingPermit := TRUE, HomingAtTargetM := btnM1, CfgHomingTargetM := 8.7, CfgTopSensorPosM := 8.7, HwIn := hw1, Cfg := cfgEncoder, Calib := calibM1); calibM1 := encoderM1.Calib;
bucketEdge(CLK := btnBucket);
encoderM2(Enable := TRUE, HomingPermit := TRUE, HomingAtTargetM := btnM2 OR bucketEdge.Q, CfgHomingTargetM := 23.7, CfgTopSensorPosM := 23.7, UseDynamicTarget := bucketEdge.Q, DynamicHomingTargetM := encoderM1.Measurement.CablePosM + cfgBucket.OffsetCloseM, HwIn := hw2, Cfg := cfgEncoder, Calib := calibM2); calibM2 := encoderM2.Calib;
bucket(Enable := TRUE, Mode := E_Mode.MAINT_N2, PowerContactorEngaged := TRUE, CablePosM1 := encoderM1.Measurement.CablePosM, CablePosM2 := encoderM2.Measurement.CablePosM, HomedM1 := encoderM1.Homed, HomedM2 := encoderM2.Homed, HomedAndReliableM1 := encoderM1.HomedAndReliable, HomedAndReliableM2 := encoderM2.HomedAndReliable, HomingSuspectM1 := encoderM1.HomingSuspect, HomingSuspectM2 := encoderM2.HomingSuspect, ConfirmClosePosition := btnBucket, Config := cfgBucket, BucketState := bucketState); bucketState := bucket.BucketState;
home.M1Status.HomedAndReliable := encoderM1.HomedAndReliable; home.M2Status.HomedAndReliable := encoderM2.HomedAndReliable; home(BucketOffsetValid := bucketState.BucketReferenced, BtnValidation := bench.Operator.JoyBtnRaw);
ADVANCE_TIME(10000000);
bench(M1_PresetTriggerCmd := encoderM1.HwOut.PresetTriggerCmd, M1_PresetValueOut := encoderM1.HwOut.PresetValueOut, M2_PresetTriggerCmd := encoderM2.HwOut.PresetTriggerCmd, M2_PresetValueOut := encoderM2.HwOut.PresetValueOut, RawPosM1 := raw1, RawPosM2 := raw2); raw1 := bench.RawPosM1; raw2 := bench.RawPosM2;
hw1.RawPosIn := bench.Winch.COD1_PosValue; hw1.SlaveOperational := TRUE; hw2.RawPosIn := bench.Winch.COD2_PosValue; hw2.SlaveOperational := TRUE;
encoderM1(Enable := TRUE, HomingPermit := TRUE, HomingAtTargetM := btnM1, CfgHomingTargetM := 8.7, CfgTopSensorPosM := 8.7, HwIn := hw1, Cfg := cfgEncoder, Calib := calibM1); calibM1 := encoderM1.Calib;
bucketEdge(CLK := btnBucket);
encoderM2(Enable := TRUE, HomingPermit := TRUE, HomingAtTargetM := btnM2 OR bucketEdge.Q, CfgHomingTargetM := 23.7, CfgTopSensorPosM := 23.7, UseDynamicTarget := bucketEdge.Q, DynamicHomingTargetM := encoderM1.Measurement.CablePosM + cfgBucket.OffsetCloseM, HwIn := hw2, Cfg := cfgEncoder, Calib := calibM2); calibM2 := encoderM2.Calib;
bucket(Enable := TRUE, Mode := E_Mode.MAINT_N2, PowerContactorEngaged := TRUE, CablePosM1 := encoderM1.Measurement.CablePosM, CablePosM2 := encoderM2.Measurement.CablePosM, HomedM1 := encoderM1.Homed, HomedM2 := encoderM2.Homed, HomedAndReliableM1 := encoderM1.HomedAndReliable, HomedAndReliableM2 := encoderM2.HomedAndReliable, HomingSuspectM1 := encoderM1.HomingSuspect, HomingSuspectM2 := encoderM2.HomingSuspect, ConfirmClosePosition := btnBucket, Config := cfgBucket, BucketState := bucketState); bucketState := bucket.BucketState;
home.M1Status.HomedAndReliable := encoderM1.HomedAndReliable; home.M2Status.HomedAndReliable := encoderM2.HomedAndReliable; home(BucketOffsetValid := bucketState.BucketReferenced, BtnValidation := bench.Operator.JoyBtnRaw);
ADVANCE_TIME(10000000);
bench(M1_PresetTriggerCmd := encoderM1.HwOut.PresetTriggerCmd, M1_PresetValueOut := encoderM1.HwOut.PresetValueOut, M2_PresetTriggerCmd := encoderM2.HwOut.PresetTriggerCmd, M2_PresetValueOut := encoderM2.HwOut.PresetValueOut, RawPosM1 := raw1, RawPosM2 := raw2); raw1 := bench.RawPosM1; raw2 := bench.RawPosM2;
hw1.RawPosIn := bench.Winch.COD1_PosValue; hw1.SlaveOperational := TRUE; hw2.RawPosIn := bench.Winch.COD2_PosValue; hw2.SlaveOperational := TRUE;
encoderM1(Enable := TRUE, HomingPermit := TRUE, HomingAtTargetM := btnM1, CfgHomingTargetM := 8.7, CfgTopSensorPosM := 8.7, HwIn := hw1, Cfg := cfgEncoder, Calib := calibM1); calibM1 := encoderM1.Calib;
bucketEdge(CLK := btnBucket);
encoderM2(Enable := TRUE, HomingPermit := TRUE, HomingAtTargetM := btnM2 OR bucketEdge.Q, CfgHomingTargetM := 23.7, CfgTopSensorPosM := 23.7, UseDynamicTarget := bucketEdge.Q, DynamicHomingTargetM := encoderM1.Measurement.CablePosM + cfgBucket.OffsetCloseM, HwIn := hw2, Cfg := cfgEncoder, Calib := calibM2); calibM2 := encoderM2.Calib;
bucket(Enable := TRUE, Mode := E_Mode.MAINT_N2, PowerContactorEngaged := TRUE, CablePosM1 := encoderM1.Measurement.CablePosM, CablePosM2 := encoderM2.Measurement.CablePosM, HomedM1 := encoderM1.Homed, HomedM2 := encoderM2.Homed, HomedAndReliableM1 := encoderM1.HomedAndReliable, HomedAndReliableM2 := encoderM2.HomedAndReliable, HomingSuspectM1 := encoderM1.HomingSuspect, HomingSuspectM2 := encoderM2.HomingSuspect, ConfirmClosePosition := btnBucket, Config := cfgBucket, BucketState := bucketState); bucketState := bucket.BucketState;
home.M1Status.HomedAndReliable := encoderM1.HomedAndReliable; home.M2Status.HomedAndReliable := encoderM2.HomedAndReliable; home(BucketOffsetValid := bucketState.BucketReferenced, BtnValidation := bench.Operator.JoyBtnRaw);
ADVANCE_TIME(10000000);
bench(M1_PresetTriggerCmd := encoderM1.HwOut.PresetTriggerCmd, M1_PresetValueOut := encoderM1.HwOut.PresetValueOut, M2_PresetTriggerCmd := encoderM2.HwOut.PresetTriggerCmd, M2_PresetValueOut := encoderM2.HwOut.PresetValueOut, RawPosM1 := raw1, RawPosM2 := raw2); raw1 := bench.RawPosM1; raw2 := bench.RawPosM2;
hw1.RawPosIn := bench.Winch.COD1_PosValue; hw1.SlaveOperational := TRUE; hw2.RawPosIn := bench.Winch.COD2_PosValue; hw2.SlaveOperational := TRUE;
encoderM1(Enable := TRUE, HomingPermit := TRUE, HomingAtTargetM := btnM1, CfgHomingTargetM := 8.7, CfgTopSensorPosM := 8.7, HwIn := hw1, Cfg := cfgEncoder, Calib := calibM1); calibM1 := encoderM1.Calib;
bucketEdge(CLK := btnBucket);
encoderM2(Enable := TRUE, HomingPermit := TRUE, HomingAtTargetM := btnM2 OR bucketEdge.Q, CfgHomingTargetM := 23.7, CfgTopSensorPosM := 23.7, UseDynamicTarget := bucketEdge.Q, DynamicHomingTargetM := encoderM1.Measurement.CablePosM + cfgBucket.OffsetCloseM, HwIn := hw2, Cfg := cfgEncoder, Calib := calibM2); calibM2 := encoderM2.Calib;
bucket(Enable := TRUE, Mode := E_Mode.MAINT_N2, PowerContactorEngaged := TRUE, CablePosM1 := encoderM1.Measurement.CablePosM, CablePosM2 := encoderM2.Measurement.CablePosM, HomedM1 := encoderM1.Homed, HomedM2 := encoderM2.Homed, HomedAndReliableM1 := encoderM1.HomedAndReliable, HomedAndReliableM2 := encoderM2.HomedAndReliable, HomingSuspectM1 := encoderM1.HomingSuspect, HomingSuspectM2 := encoderM2.HomingSuspect, ConfirmClosePosition := btnBucket, Config := cfgBucket, BucketState := bucketState); bucketState := bucket.BucketState;
home.M1Status.HomedAndReliable := encoderM1.HomedAndReliable; home.M2Status.HomedAndReliable := encoderM2.HomedAndReliable; home(BucketOffsetValid := bucketState.BucketReferenced, BtnValidation := bench.Operator.JoyBtnRaw);
ADVANCE_TIME(10000000);
bench(M1_PresetTriggerCmd := encoderM1.HwOut.PresetTriggerCmd, M1_PresetValueOut := encoderM1.HwOut.PresetValueOut, M2_PresetTriggerCmd := encoderM2.HwOut.PresetTriggerCmd, M2_PresetValueOut := encoderM2.HwOut.PresetValueOut, RawPosM1 := raw1, RawPosM2 := raw2); raw1 := bench.RawPosM1; raw2 := bench.RawPosM2;
hw1.RawPosIn := bench.Winch.COD1_PosValue; hw1.SlaveOperational := TRUE; hw2.RawPosIn := bench.Winch.COD2_PosValue; hw2.SlaveOperational := TRUE;
encoderM1(Enable := TRUE, HomingPermit := TRUE, HomingAtTargetM := btnM1, CfgHomingTargetM := 8.7, CfgTopSensorPosM := 8.7, HwIn := hw1, Cfg := cfgEncoder, Calib := calibM1); calibM1 := encoderM1.Calib;
bucketEdge(CLK := btnBucket);
encoderM2(Enable := TRUE, HomingPermit := TRUE, HomingAtTargetM := btnM2 OR bucketEdge.Q, CfgHomingTargetM := 23.7, CfgTopSensorPosM := 23.7, UseDynamicTarget := bucketEdge.Q, DynamicHomingTargetM := encoderM1.Measurement.CablePosM + cfgBucket.OffsetCloseM, HwIn := hw2, Cfg := cfgEncoder, Calib := calibM2); calibM2 := encoderM2.Calib;
bucket(Enable := TRUE, Mode := E_Mode.MAINT_N2, PowerContactorEngaged := TRUE, CablePosM1 := encoderM1.Measurement.CablePosM, CablePosM2 := encoderM2.Measurement.CablePosM, HomedM1 := encoderM1.Homed, HomedM2 := encoderM2.Homed, HomedAndReliableM1 := encoderM1.HomedAndReliable, HomedAndReliableM2 := encoderM2.HomedAndReliable, HomingSuspectM1 := encoderM1.HomingSuspect, HomingSuspectM2 := encoderM2.HomingSuspect, ConfirmClosePosition := btnBucket, Config := cfgBucket, BucketState := bucketState); bucketState := bucket.BucketState;
home.M1Status.HomedAndReliable := encoderM1.HomedAndReliable; home.M2Status.HomedAndReliable := encoderM2.HomedAndReliable; home(BucketOffsetValid := bucketState.BucketReferenced, BtnValidation := bench.Operator.JoyBtnRaw);
ADVANCE_TIME(10000000);
bench(M1_PresetTriggerCmd := encoderM1.HwOut.PresetTriggerCmd, M1_PresetValueOut := encoderM1.HwOut.PresetValueOut, M2_PresetTriggerCmd := encoderM2.HwOut.PresetTriggerCmd, M2_PresetValueOut := encoderM2.HwOut.PresetValueOut, RawPosM1 := raw1, RawPosM2 := raw2); raw1 := bench.RawPosM1; raw2 := bench.RawPosM2;
hw1.RawPosIn := bench.Winch.COD1_PosValue; hw1.SlaveOperational := TRUE; hw2.RawPosIn := bench.Winch.COD2_PosValue; hw2.SlaveOperational := TRUE;
encoderM1(Enable := TRUE, HomingPermit := TRUE, HomingAtTargetM := btnM1, CfgHomingTargetM := 8.7, CfgTopSensorPosM := 8.7, HwIn := hw1, Cfg := cfgEncoder, Calib := calibM1); calibM1 := encoderM1.Calib;
bucketEdge(CLK := btnBucket);
encoderM2(Enable := TRUE, HomingPermit := TRUE, HomingAtTargetM := btnM2 OR bucketEdge.Q, CfgHomingTargetM := 23.7, CfgTopSensorPosM := 23.7, UseDynamicTarget := bucketEdge.Q, DynamicHomingTargetM := encoderM1.Measurement.CablePosM + cfgBucket.OffsetCloseM, HwIn := hw2, Cfg := cfgEncoder, Calib := calibM2); calibM2 := encoderM2.Calib;
bucket(Enable := TRUE, Mode := E_Mode.MAINT_N2, PowerContactorEngaged := TRUE, CablePosM1 := encoderM1.Measurement.CablePosM, CablePosM2 := encoderM2.Measurement.CablePosM, HomedM1 := encoderM1.Homed, HomedM2 := encoderM2.Homed, HomedAndReliableM1 := encoderM1.HomedAndReliable, HomedAndReliableM2 := encoderM2.HomedAndReliable, HomingSuspectM1 := encoderM1.HomingSuspect, HomingSuspectM2 := encoderM2.HomingSuspect, ConfirmClosePosition := btnBucket, Config := cfgBucket, BucketState := bucketState); bucketState := bucket.BucketState;
home.M1Status.HomedAndReliable := encoderM1.HomedAndReliable; home.M2Status.HomedAndReliable := encoderM2.HomedAndReliable; home(BucketOffsetValid := bucketState.BucketReferenced, BtnValidation := bench.Operator.JoyBtnRaw);
ADVANCE_TIME(10000000);
bench(M1_PresetTriggerCmd := encoderM1.HwOut.PresetTriggerCmd, M1_PresetValueOut := encoderM1.HwOut.PresetValueOut, M2_PresetTriggerCmd := encoderM2.HwOut.PresetTriggerCmd, M2_PresetValueOut := encoderM2.HwOut.PresetValueOut, RawPosM1 := raw1, RawPosM2 := raw2); raw1 := bench.RawPosM1; raw2 := bench.RawPosM2;
hw1.RawPosIn := bench.Winch.COD1_PosValue; hw1.SlaveOperational := TRUE; hw2.RawPosIn := bench.Winch.COD2_PosValue; hw2.SlaveOperational := TRUE;
encoderM1(Enable := TRUE, HomingPermit := TRUE, HomingAtTargetM := btnM1, CfgHomingTargetM := 8.7, CfgTopSensorPosM := 8.7, HwIn := hw1, Cfg := cfgEncoder, Calib := calibM1); calibM1 := encoderM1.Calib;
bucketEdge(CLK := btnBucket);
encoderM2(Enable := TRUE, HomingPermit := TRUE, HomingAtTargetM := btnM2 OR bucketEdge.Q, CfgHomingTargetM := 23.7, CfgTopSensorPosM := 23.7, UseDynamicTarget := bucketEdge.Q, DynamicHomingTargetM := encoderM1.Measurement.CablePosM + cfgBucket.OffsetCloseM, HwIn := hw2, Cfg := cfgEncoder, Calib := calibM2); calibM2 := encoderM2.Calib;
bucket(Enable := TRUE, Mode := E_Mode.MAINT_N2, PowerContactorEngaged := TRUE, CablePosM1 := encoderM1.Measurement.CablePosM, CablePosM2 := encoderM2.Measurement.CablePosM, HomedM1 := encoderM1.Homed, HomedM2 := encoderM2.Homed, HomedAndReliableM1 := encoderM1.HomedAndReliable, HomedAndReliableM2 := encoderM2.HomedAndReliable, HomingSuspectM1 := encoderM1.HomingSuspect, HomingSuspectM2 := encoderM2.HomingSuspect, ConfirmClosePosition := btnBucket, Config := cfgBucket, BucketState := bucketState); bucketState := bucket.BucketState;
home.M1Status.HomedAndReliable := encoderM1.HomedAndReliable; home.M2Status.HomedAndReliable := encoderM2.HomedAndReliable; home(BucketOffsetValid := bucketState.BucketReferenced, BtnValidation := bench.Operator.JoyBtnRaw);
ADVANCE_TIME(10000000);
bench(M1_PresetTriggerCmd := encoderM1.HwOut.PresetTriggerCmd, M1_PresetValueOut := encoderM1.HwOut.PresetValueOut, M2_PresetTriggerCmd := encoderM2.HwOut.PresetTriggerCmd, M2_PresetValueOut := encoderM2.HwOut.PresetValueOut, RawPosM1 := raw1, RawPosM2 := raw2); raw1 := bench.RawPosM1; raw2 := bench.RawPosM2;
hw1.RawPosIn := bench.Winch.COD1_PosValue; hw1.SlaveOperational := TRUE; hw2.RawPosIn := bench.Winch.COD2_PosValue; hw2.SlaveOperational := TRUE;
encoderM1(Enable := TRUE, HomingPermit := TRUE, HomingAtTargetM := btnM1, CfgHomingTargetM := 8.7, CfgTopSensorPosM := 8.7, HwIn := hw1, Cfg := cfgEncoder, Calib := calibM1); calibM1 := encoderM1.Calib;
bucketEdge(CLK := btnBucket);
encoderM2(Enable := TRUE, HomingPermit := TRUE, HomingAtTargetM := btnM2 OR bucketEdge.Q, CfgHomingTargetM := 23.7, CfgTopSensorPosM := 23.7, UseDynamicTarget := bucketEdge.Q, DynamicHomingTargetM := encoderM1.Measurement.CablePosM + cfgBucket.OffsetCloseM, HwIn := hw2, Cfg := cfgEncoder, Calib := calibM2); calibM2 := encoderM2.Calib;
bucket(Enable := TRUE, Mode := E_Mode.MAINT_N2, PowerContactorEngaged := TRUE, CablePosM1 := encoderM1.Measurement.CablePosM, CablePosM2 := encoderM2.Measurement.CablePosM, HomedM1 := encoderM1.Homed, HomedM2 := encoderM2.Homed, HomedAndReliableM1 := encoderM1.HomedAndReliable, HomedAndReliableM2 := encoderM2.HomedAndReliable, HomingSuspectM1 := encoderM1.HomingSuspect, HomingSuspectM2 := encoderM2.HomingSuspect, ConfirmClosePosition := btnBucket, Config := cfgBucket, BucketState := bucketState); bucketState := bucket.BucketState;
home.M1Status.HomedAndReliable := encoderM1.HomedAndReliable; home.M2Status.HomedAndReliable := encoderM2.HomedAndReliable; home(BucketOffsetValid := bucketState.BucketReferenced, BtnValidation := bench.Operator.JoyBtnRaw);
ADVANCE_TIME(10000000);
bench(M1_PresetTriggerCmd := encoderM1.HwOut.PresetTriggerCmd, M1_PresetValueOut := encoderM1.HwOut.PresetValueOut, M2_PresetTriggerCmd := encoderM2.HwOut.PresetTriggerCmd, M2_PresetValueOut := encoderM2.HwOut.PresetValueOut, RawPosM1 := raw1, RawPosM2 := raw2); raw1 := bench.RawPosM1; raw2 := bench.RawPosM2;
hw1.RawPosIn := bench.Winch.COD1_PosValue; hw1.SlaveOperational := TRUE; hw2.RawPosIn := bench.Winch.COD2_PosValue; hw2.SlaveOperational := TRUE;
encoderM1(Enable := TRUE, HomingPermit := TRUE, HomingAtTargetM := btnM1, CfgHomingTargetM := 8.7, CfgTopSensorPosM := 8.7, HwIn := hw1, Cfg := cfgEncoder, Calib := calibM1); calibM1 := encoderM1.Calib;
bucketEdge(CLK := btnBucket);
encoderM2(Enable := TRUE, HomingPermit := TRUE, HomingAtTargetM := btnM2 OR bucketEdge.Q, CfgHomingTargetM := 23.7, CfgTopSensorPosM := 23.7, UseDynamicTarget := bucketEdge.Q, DynamicHomingTargetM := encoderM1.Measurement.CablePosM + cfgBucket.OffsetCloseM, HwIn := hw2, Cfg := cfgEncoder, Calib := calibM2); calibM2 := encoderM2.Calib;
bucket(Enable := TRUE, Mode := E_Mode.MAINT_N2, PowerContactorEngaged := TRUE, CablePosM1 := encoderM1.Measurement.CablePosM, CablePosM2 := encoderM2.Measurement.CablePosM, HomedM1 := encoderM1.Homed, HomedM2 := encoderM2.Homed, HomedAndReliableM1 := encoderM1.HomedAndReliable, HomedAndReliableM2 := encoderM2.HomedAndReliable, HomingSuspectM1 := encoderM1.HomingSuspect, HomingSuspectM2 := encoderM2.HomingSuspect, ConfirmClosePosition := btnBucket, Config := cfgBucket, BucketState := bucketState); bucketState := bucket.BucketState;
home.M1Status.HomedAndReliable := encoderM1.HomedAndReliable; home.M2Status.HomedAndReliable := encoderM2.HomedAndReliable; home(BucketOffsetValid := bucketState.BucketReferenced, BtnValidation := bench.Operator.JoyBtnRaw);
ADVANCE_TIME(10000000);
bench(M1_PresetTriggerCmd := encoderM1.HwOut.PresetTriggerCmd, M1_PresetValueOut := encoderM1.HwOut.PresetValueOut, M2_PresetTriggerCmd := encoderM2.HwOut.PresetTriggerCmd, M2_PresetValueOut := encoderM2.HwOut.PresetValueOut, RawPosM1 := raw1, RawPosM2 := raw2); raw1 := bench.RawPosM1; raw2 := bench.RawPosM2;
hw1.RawPosIn := bench.Winch.COD1_PosValue; hw1.SlaveOperational := TRUE; hw2.RawPosIn := bench.Winch.COD2_PosValue; hw2.SlaveOperational := TRUE;
encoderM1(Enable := TRUE, HomingPermit := TRUE, HomingAtTargetM := btnM1, CfgHomingTargetM := 8.7, CfgTopSensorPosM := 8.7, HwIn := hw1, Cfg := cfgEncoder, Calib := calibM1); calibM1 := encoderM1.Calib;
bucketEdge(CLK := btnBucket);
encoderM2(Enable := TRUE, HomingPermit := TRUE, HomingAtTargetM := btnM2 OR bucketEdge.Q, CfgHomingTargetM := 23.7, CfgTopSensorPosM := 23.7, UseDynamicTarget := bucketEdge.Q, DynamicHomingTargetM := encoderM1.Measurement.CablePosM + cfgBucket.OffsetCloseM, HwIn := hw2, Cfg := cfgEncoder, Calib := calibM2); calibM2 := encoderM2.Calib;
bucket(Enable := TRUE, Mode := E_Mode.MAINT_N2, PowerContactorEngaged := TRUE, CablePosM1 := encoderM1.Measurement.CablePosM, CablePosM2 := encoderM2.Measurement.CablePosM, HomedM1 := encoderM1.Homed, HomedM2 := encoderM2.Homed, HomedAndReliableM1 := encoderM1.HomedAndReliable, HomedAndReliableM2 := encoderM2.HomedAndReliable, HomingSuspectM1 := encoderM1.HomingSuspect, HomingSuspectM2 := encoderM2.HomingSuspect, ConfirmClosePosition := btnBucket, Config := cfgBucket, BucketState := bucketState); bucketState := bucket.BucketState;
home.M1Status.HomedAndReliable := encoderM1.HomedAndReliable; home.M2Status.HomedAndReliable := encoderM2.HomedAndReliable; home(BucketOffsetValid := bucketState.BucketReferenced, BtnValidation := bench.Operator.JoyBtnRaw);
ADVANCE_TIME(10000000);
bench(M1_PresetTriggerCmd := encoderM1.HwOut.PresetTriggerCmd, M1_PresetValueOut := encoderM1.HwOut.PresetValueOut, M2_PresetTriggerCmd := encoderM2.HwOut.PresetTriggerCmd, M2_PresetValueOut := encoderM2.HwOut.PresetValueOut, RawPosM1 := raw1, RawPosM2 := raw2); raw1 := bench.RawPosM1; raw2 := bench.RawPosM2;
hw1.RawPosIn := bench.Winch.COD1_PosValue; hw1.SlaveOperational := TRUE; hw2.RawPosIn := bench.Winch.COD2_PosValue; hw2.SlaveOperational := TRUE;
encoderM1(Enable := TRUE, HomingPermit := TRUE, HomingAtTargetM := btnM1, CfgHomingTargetM := 8.7, CfgTopSensorPosM := 8.7, HwIn := hw1, Cfg := cfgEncoder, Calib := calibM1); calibM1 := encoderM1.Calib;
bucketEdge(CLK := btnBucket);
encoderM2(Enable := TRUE, HomingPermit := TRUE, HomingAtTargetM := btnM2 OR bucketEdge.Q, CfgHomingTargetM := 23.7, CfgTopSensorPosM := 23.7, UseDynamicTarget := bucketEdge.Q, DynamicHomingTargetM := encoderM1.Measurement.CablePosM + cfgBucket.OffsetCloseM, HwIn := hw2, Cfg := cfgEncoder, Calib := calibM2); calibM2 := encoderM2.Calib;
bucket(Enable := TRUE, Mode := E_Mode.MAINT_N2, PowerContactorEngaged := TRUE, CablePosM1 := encoderM1.Measurement.CablePosM, CablePosM2 := encoderM2.Measurement.CablePosM, HomedM1 := encoderM1.Homed, HomedM2 := encoderM2.Homed, HomedAndReliableM1 := encoderM1.HomedAndReliable, HomedAndReliableM2 := encoderM2.HomedAndReliable, HomingSuspectM1 := encoderM1.HomingSuspect, HomingSuspectM2 := encoderM2.HomingSuspect, ConfirmClosePosition := btnBucket, Config := cfgBucket, BucketState := bucketState); bucketState := bucket.BucketState;
home.M1Status.HomedAndReliable := encoderM1.HomedAndReliable; home.M2Status.HomedAndReliable := encoderM2.HomedAndReliable; home(BucketOffsetValid := bucketState.BucketReferenced, BtnValidation := bench.Operator.JoyBtnRaw);
ADVANCE_TIME(10000000);
bench(M1_PresetTriggerCmd := encoderM1.HwOut.PresetTriggerCmd, M1_PresetValueOut := encoderM1.HwOut.PresetValueOut, M2_PresetTriggerCmd := encoderM2.HwOut.PresetTriggerCmd, M2_PresetValueOut := encoderM2.HwOut.PresetValueOut, RawPosM1 := raw1, RawPosM2 := raw2); raw1 := bench.RawPosM1; raw2 := bench.RawPosM2;
hw1.RawPosIn := bench.Winch.COD1_PosValue; hw1.SlaveOperational := TRUE; hw2.RawPosIn := bench.Winch.COD2_PosValue; hw2.SlaveOperational := TRUE;
encoderM1(Enable := TRUE, HomingPermit := TRUE, HomingAtTargetM := btnM1, CfgHomingTargetM := 8.7, CfgTopSensorPosM := 8.7, HwIn := hw1, Cfg := cfgEncoder, Calib := calibM1); calibM1 := encoderM1.Calib;
bucketEdge(CLK := btnBucket);
encoderM2(Enable := TRUE, HomingPermit := TRUE, HomingAtTargetM := btnM2 OR bucketEdge.Q, CfgHomingTargetM := 23.7, CfgTopSensorPosM := 23.7, UseDynamicTarget := bucketEdge.Q, DynamicHomingTargetM := encoderM1.Measurement.CablePosM + cfgBucket.OffsetCloseM, HwIn := hw2, Cfg := cfgEncoder, Calib := calibM2); calibM2 := encoderM2.Calib;
bucket(Enable := TRUE, Mode := E_Mode.MAINT_N2, PowerContactorEngaged := TRUE, CablePosM1 := encoderM1.Measurement.CablePosM, CablePosM2 := encoderM2.Measurement.CablePosM, HomedM1 := encoderM1.Homed, HomedM2 := encoderM2.Homed, HomedAndReliableM1 := encoderM1.HomedAndReliable, HomedAndReliableM2 := encoderM2.HomedAndReliable, HomingSuspectM1 := encoderM1.HomingSuspect, HomingSuspectM2 := encoderM2.HomingSuspect, ConfirmClosePosition := btnBucket, Config := cfgBucket, BucketState := bucketState); bucketState := bucket.BucketState;
home.M1Status.HomedAndReliable := encoderM1.HomedAndReliable; home.M2Status.HomedAndReliable := encoderM2.HomedAndReliable; home(BucketOffsetValid := bucketState.BucketReferenced, BtnValidation := bench.Operator.JoyBtnRaw);
ADVANCE_TIME(10000000);
bench(M1_PresetTriggerCmd := encoderM1.HwOut.PresetTriggerCmd, M1_PresetValueOut := encoderM1.HwOut.PresetValueOut, M2_PresetTriggerCmd := encoderM2.HwOut.PresetTriggerCmd, M2_PresetValueOut := encoderM2.HwOut.PresetValueOut, RawPosM1 := raw1, RawPosM2 := raw2); raw1 := bench.RawPosM1; raw2 := bench.RawPosM2;
hw1.RawPosIn := bench.Winch.COD1_PosValue; hw1.SlaveOperational := TRUE; hw2.RawPosIn := bench.Winch.COD2_PosValue; hw2.SlaveOperational := TRUE;
encoderM1(Enable := TRUE, HomingPermit := TRUE, HomingAtTargetM := btnM1, CfgHomingTargetM := 8.7, CfgTopSensorPosM := 8.7, HwIn := hw1, Cfg := cfgEncoder, Calib := calibM1); calibM1 := encoderM1.Calib;
bucketEdge(CLK := btnBucket);
encoderM2(Enable := TRUE, HomingPermit := TRUE, HomingAtTargetM := btnM2 OR bucketEdge.Q, CfgHomingTargetM := 23.7, CfgTopSensorPosM := 23.7, UseDynamicTarget := bucketEdge.Q, DynamicHomingTargetM := encoderM1.Measurement.CablePosM + cfgBucket.OffsetCloseM, HwIn := hw2, Cfg := cfgEncoder, Calib := calibM2); calibM2 := encoderM2.Calib;
bucket(Enable := TRUE, Mode := E_Mode.MAINT_N2, PowerContactorEngaged := TRUE, CablePosM1 := encoderM1.Measurement.CablePosM, CablePosM2 := encoderM2.Measurement.CablePosM, HomedM1 := encoderM1.Homed, HomedM2 := encoderM2.Homed, HomedAndReliableM1 := encoderM1.HomedAndReliable, HomedAndReliableM2 := encoderM2.HomedAndReliable, HomingSuspectM1 := encoderM1.HomingSuspect, HomingSuspectM2 := encoderM2.HomingSuspect, ConfirmClosePosition := btnBucket, Config := cfgBucket, BucketState := bucketState); bucketState := bucket.BucketState;
home.M1Status.HomedAndReliable := encoderM1.HomedAndReliable; home.M2Status.HomedAndReliable := encoderM2.HomedAndReliable; home(BucketOffsetValid := bucketState.BucketReferenced, BtnValidation := bench.Operator.JoyBtnRaw);
ADVANCE_TIME(10000000);
bench(M1_PresetTriggerCmd := encoderM1.HwOut.PresetTriggerCmd, M1_PresetValueOut := encoderM1.HwOut.PresetValueOut, M2_PresetTriggerCmd := encoderM2.HwOut.PresetTriggerCmd, M2_PresetValueOut := encoderM2.HwOut.PresetValueOut, RawPosM1 := raw1, RawPosM2 := raw2); raw1 := bench.RawPosM1; raw2 := bench.RawPosM2;
hw1.RawPosIn := bench.Winch.COD1_PosValue; hw1.SlaveOperational := TRUE; hw2.RawPosIn := bench.Winch.COD2_PosValue; hw2.SlaveOperational := TRUE;
encoderM1(Enable := TRUE, HomingPermit := TRUE, HomingAtTargetM := btnM1, CfgHomingTargetM := 8.7, CfgTopSensorPosM := 8.7, HwIn := hw1, Cfg := cfgEncoder, Calib := calibM1); calibM1 := encoderM1.Calib;
bucketEdge(CLK := btnBucket);
encoderM2(Enable := TRUE, HomingPermit := TRUE, HomingAtTargetM := btnM2 OR bucketEdge.Q, CfgHomingTargetM := 23.7, CfgTopSensorPosM := 23.7, UseDynamicTarget := bucketEdge.Q, DynamicHomingTargetM := encoderM1.Measurement.CablePosM + cfgBucket.OffsetCloseM, HwIn := hw2, Cfg := cfgEncoder, Calib := calibM2); calibM2 := encoderM2.Calib;
bucket(Enable := TRUE, Mode := E_Mode.MAINT_N2, PowerContactorEngaged := TRUE, CablePosM1 := encoderM1.Measurement.CablePosM, CablePosM2 := encoderM2.Measurement.CablePosM, HomedM1 := encoderM1.Homed, HomedM2 := encoderM2.Homed, HomedAndReliableM1 := encoderM1.HomedAndReliable, HomedAndReliableM2 := encoderM2.HomedAndReliable, HomingSuspectM1 := encoderM1.HomingSuspect, HomingSuspectM2 := encoderM2.HomingSuspect, ConfirmClosePosition := btnBucket, Config := cfgBucket, BucketState := bucketState); bucketState := bucket.BucketState;
home.M1Status.HomedAndReliable := encoderM1.HomedAndReliable; home.M2Status.HomedAndReliable := encoderM2.HomedAndReliable; home(BucketOffsetValid := bucketState.BucketReferenced, BtnValidation := bench.Operator.JoyBtnRaw);
ADVANCE_TIME(10000000);
bench(M1_PresetTriggerCmd := encoderM1.HwOut.PresetTriggerCmd, M1_PresetValueOut := encoderM1.HwOut.PresetValueOut, M2_PresetTriggerCmd := encoderM2.HwOut.PresetTriggerCmd, M2_PresetValueOut := encoderM2.HwOut.PresetValueOut, RawPosM1 := raw1, RawPosM2 := raw2); raw1 := bench.RawPosM1; raw2 := bench.RawPosM2;
hw1.RawPosIn := bench.Winch.COD1_PosValue; hw1.SlaveOperational := TRUE; hw2.RawPosIn := bench.Winch.COD2_PosValue; hw2.SlaveOperational := TRUE;
encoderM1(Enable := TRUE, HomingPermit := TRUE, HomingAtTargetM := btnM1, CfgHomingTargetM := 8.7, CfgTopSensorPosM := 8.7, HwIn := hw1, Cfg := cfgEncoder, Calib := calibM1); calibM1 := encoderM1.Calib;
bucketEdge(CLK := btnBucket);
encoderM2(Enable := TRUE, HomingPermit := TRUE, HomingAtTargetM := btnM2 OR bucketEdge.Q, CfgHomingTargetM := 23.7, CfgTopSensorPosM := 23.7, UseDynamicTarget := bucketEdge.Q, DynamicHomingTargetM := encoderM1.Measurement.CablePosM + cfgBucket.OffsetCloseM, HwIn := hw2, Cfg := cfgEncoder, Calib := calibM2); calibM2 := encoderM2.Calib;
bucket(Enable := TRUE, Mode := E_Mode.MAINT_N2, PowerContactorEngaged := TRUE, CablePosM1 := encoderM1.Measurement.CablePosM, CablePosM2 := encoderM2.Measurement.CablePosM, HomedM1 := encoderM1.Homed, HomedM2 := encoderM2.Homed, HomedAndReliableM1 := encoderM1.HomedAndReliable, HomedAndReliableM2 := encoderM2.HomedAndReliable, HomingSuspectM1 := encoderM1.HomingSuspect, HomingSuspectM2 := encoderM2.HomingSuspect, ConfirmClosePosition := btnBucket, Config := cfgBucket, BucketState := bucketState); bucketState := bucket.BucketState;
home.M1Status.HomedAndReliable := encoderM1.HomedAndReliable; home.M2Status.HomedAndReliable := encoderM2.HomedAndReliable; home(BucketOffsetValid := bucketState.BucketReferenced, BtnValidation := bench.Operator.JoyBtnRaw);
ADVANCE_TIME(10000000);
bench(M1_PresetTriggerCmd := encoderM1.HwOut.PresetTriggerCmd, M1_PresetValueOut := encoderM1.HwOut.PresetValueOut, M2_PresetTriggerCmd := encoderM2.HwOut.PresetTriggerCmd, M2_PresetValueOut := encoderM2.HwOut.PresetValueOut, RawPosM1 := raw1, RawPosM2 := raw2); raw1 := bench.RawPosM1; raw2 := bench.RawPosM2;
hw1.RawPosIn := bench.Winch.COD1_PosValue; hw1.SlaveOperational := TRUE; hw2.RawPosIn := bench.Winch.COD2_PosValue; hw2.SlaveOperational := TRUE;
encoderM1(Enable := TRUE, HomingPermit := TRUE, HomingAtTargetM := btnM1, CfgHomingTargetM := 8.7, CfgTopSensorPosM := 8.7, HwIn := hw1, Cfg := cfgEncoder, Calib := calibM1); calibM1 := encoderM1.Calib;
bucketEdge(CLK := btnBucket);
encoderM2(Enable := TRUE, HomingPermit := TRUE, HomingAtTargetM := btnM2 OR bucketEdge.Q, CfgHomingTargetM := 23.7, CfgTopSensorPosM := 23.7, UseDynamicTarget := bucketEdge.Q, DynamicHomingTargetM := encoderM1.Measurement.CablePosM + cfgBucket.OffsetCloseM, HwIn := hw2, Cfg := cfgEncoder, Calib := calibM2); calibM2 := encoderM2.Calib;
bucket(Enable := TRUE, Mode := E_Mode.MAINT_N2, PowerContactorEngaged := TRUE, CablePosM1 := encoderM1.Measurement.CablePosM, CablePosM2 := encoderM2.Measurement.CablePosM, HomedM1 := encoderM1.Homed, HomedM2 := encoderM2.Homed, HomedAndReliableM1 := encoderM1.HomedAndReliable, HomedAndReliableM2 := encoderM2.HomedAndReliable, HomingSuspectM1 := encoderM1.HomingSuspect, HomingSuspectM2 := encoderM2.HomingSuspect, ConfirmClosePosition := btnBucket, Config := cfgBucket, BucketState := bucketState); bucketState := bucket.BucketState;
home.M1Status.HomedAndReliable := encoderM1.HomedAndReliable; home.M2Status.HomedAndReliable := encoderM2.HomedAndReliable; home(BucketOffsetValid := bucketState.BucketReferenced, BtnValidation := bench.Operator.JoyBtnRaw);
ADVANCE_TIME(10000000);
bench(M1_PresetTriggerCmd := encoderM1.HwOut.PresetTriggerCmd, M1_PresetValueOut := encoderM1.HwOut.PresetValueOut, M2_PresetTriggerCmd := encoderM2.HwOut.PresetTriggerCmd, M2_PresetValueOut := encoderM2.HwOut.PresetValueOut, RawPosM1 := raw1, RawPosM2 := raw2); raw1 := bench.RawPosM1; raw2 := bench.RawPosM2;
hw1.RawPosIn := bench.Winch.COD1_PosValue; hw1.SlaveOperational := TRUE; hw2.RawPosIn := bench.Winch.COD2_PosValue; hw2.SlaveOperational := TRUE;
encoderM1(Enable := TRUE, HomingPermit := TRUE, HomingAtTargetM := btnM1, CfgHomingTargetM := 8.7, CfgTopSensorPosM := 8.7, HwIn := hw1, Cfg := cfgEncoder, Calib := calibM1); calibM1 := encoderM1.Calib;
bucketEdge(CLK := btnBucket);
encoderM2(Enable := TRUE, HomingPermit := TRUE, HomingAtTargetM := btnM2 OR bucketEdge.Q, CfgHomingTargetM := 23.7, CfgTopSensorPosM := 23.7, UseDynamicTarget := bucketEdge.Q, DynamicHomingTargetM := encoderM1.Measurement.CablePosM + cfgBucket.OffsetCloseM, HwIn := hw2, Cfg := cfgEncoder, Calib := calibM2); calibM2 := encoderM2.Calib;
bucket(Enable := TRUE, Mode := E_Mode.MAINT_N2, PowerContactorEngaged := TRUE, CablePosM1 := encoderM1.Measurement.CablePosM, CablePosM2 := encoderM2.Measurement.CablePosM, HomedM1 := encoderM1.Homed, HomedM2 := encoderM2.Homed, HomedAndReliableM1 := encoderM1.HomedAndReliable, HomedAndReliableM2 := encoderM2.HomedAndReliable, HomingSuspectM1 := encoderM1.HomingSuspect, HomingSuspectM2 := encoderM2.HomingSuspect, ConfirmClosePosition := btnBucket, Config := cfgBucket, BucketState := bucketState); bucketState := bucket.BucketState;
home.M1Status.HomedAndReliable := encoderM1.HomedAndReliable; home.M2Status.HomedAndReliable := encoderM2.HomedAndReliable; home(BucketOffsetValid := bucketState.BucketReferenced, BtnValidation := bench.Operator.JoyBtnRaw);
ADVANCE_TIME(10000000);
bench(M1_PresetTriggerCmd := encoderM1.HwOut.PresetTriggerCmd, M1_PresetValueOut := encoderM1.HwOut.PresetValueOut, M2_PresetTriggerCmd := encoderM2.HwOut.PresetTriggerCmd, M2_PresetValueOut := encoderM2.HwOut.PresetValueOut, RawPosM1 := raw1, RawPosM2 := raw2); raw1 := bench.RawPosM1; raw2 := bench.RawPosM2;
hw1.RawPosIn := bench.Winch.COD1_PosValue; hw1.SlaveOperational := TRUE; hw2.RawPosIn := bench.Winch.COD2_PosValue; hw2.SlaveOperational := TRUE;
encoderM1(Enable := TRUE, HomingPermit := TRUE, HomingAtTargetM := btnM1, CfgHomingTargetM := 8.7, CfgTopSensorPosM := 8.7, HwIn := hw1, Cfg := cfgEncoder, Calib := calibM1); calibM1 := encoderM1.Calib;
bucketEdge(CLK := btnBucket);
encoderM2(Enable := TRUE, HomingPermit := TRUE, HomingAtTargetM := btnM2 OR bucketEdge.Q, CfgHomingTargetM := 23.7, CfgTopSensorPosM := 23.7, UseDynamicTarget := bucketEdge.Q, DynamicHomingTargetM := encoderM1.Measurement.CablePosM + cfgBucket.OffsetCloseM, HwIn := hw2, Cfg := cfgEncoder, Calib := calibM2); calibM2 := encoderM2.Calib;
bucket(Enable := TRUE, Mode := E_Mode.MAINT_N2, PowerContactorEngaged := TRUE, CablePosM1 := encoderM1.Measurement.CablePosM, CablePosM2 := encoderM2.Measurement.CablePosM, HomedM1 := encoderM1.Homed, HomedM2 := encoderM2.Homed, HomedAndReliableM1 := encoderM1.HomedAndReliable, HomedAndReliableM2 := encoderM2.HomedAndReliable, HomingSuspectM1 := encoderM1.HomingSuspect, HomingSuspectM2 := encoderM2.HomingSuspect, ConfirmClosePosition := btnBucket, Config := cfgBucket, BucketState := bucketState); bucketState := bucket.BucketState;
home.M1Status.HomedAndReliable := encoderM1.HomedAndReliable; home.M2Status.HomedAndReliable := encoderM2.HomedAndReliable; home(BucketOffsetValid := bucketState.BucketReferenced, BtnValidation := bench.Operator.JoyBtnRaw);
ADVANCE_TIME(10000000);
bench(M1_PresetTriggerCmd := encoderM1.HwOut.PresetTriggerCmd, M1_PresetValueOut := encoderM1.HwOut.PresetValueOut, M2_PresetTriggerCmd := encoderM2.HwOut.PresetTriggerCmd, M2_PresetValueOut := encoderM2.HwOut.PresetValueOut, RawPosM1 := raw1, RawPosM2 := raw2); raw1 := bench.RawPosM1; raw2 := bench.RawPosM2;
hw1.RawPosIn := bench.Winch.COD1_PosValue; hw1.SlaveOperational := TRUE; hw2.RawPosIn := bench.Winch.COD2_PosValue; hw2.SlaveOperational := TRUE;
encoderM1(Enable := TRUE, HomingPermit := TRUE, HomingAtTargetM := btnM1, CfgHomingTargetM := 8.7, CfgTopSensorPosM := 8.7, HwIn := hw1, Cfg := cfgEncoder, Calib := calibM1); calibM1 := encoderM1.Calib;
bucketEdge(CLK := btnBucket);
encoderM2(Enable := TRUE, HomingPermit := TRUE, HomingAtTargetM := btnM2 OR bucketEdge.Q, CfgHomingTargetM := 23.7, CfgTopSensorPosM := 23.7, UseDynamicTarget := bucketEdge.Q, DynamicHomingTargetM := encoderM1.Measurement.CablePosM + cfgBucket.OffsetCloseM, HwIn := hw2, Cfg := cfgEncoder, Calib := calibM2); calibM2 := encoderM2.Calib;
bucket(Enable := TRUE, Mode := E_Mode.MAINT_N2, PowerContactorEngaged := TRUE, CablePosM1 := encoderM1.Measurement.CablePosM, CablePosM2 := encoderM2.Measurement.CablePosM, HomedM1 := encoderM1.Homed, HomedM2 := encoderM2.Homed, HomedAndReliableM1 := encoderM1.HomedAndReliable, HomedAndReliableM2 := encoderM2.HomedAndReliable, HomingSuspectM1 := encoderM1.HomingSuspect, HomingSuspectM2 := encoderM2.HomingSuspect, ConfirmClosePosition := btnBucket, Config := cfgBucket, BucketState := bucketState); bucketState := bucket.BucketState;
home.M1Status.HomedAndReliable := encoderM1.HomedAndReliable; home.M2Status.HomedAndReliable := encoderM2.HomedAndReliable; home(BucketOffsetValid := bucketState.BucketReferenced, BtnValidation := bench.Operator.JoyBtnRaw);
ADVANCE_TIME(10000000);
bench(M1_PresetTriggerCmd := encoderM1.HwOut.PresetTriggerCmd, M1_PresetValueOut := encoderM1.HwOut.PresetValueOut, M2_PresetTriggerCmd := encoderM2.HwOut.PresetTriggerCmd, M2_PresetValueOut := encoderM2.HwOut.PresetValueOut, RawPosM1 := raw1, RawPosM2 := raw2); raw1 := bench.RawPosM1; raw2 := bench.RawPosM2;
hw1.RawPosIn := bench.Winch.COD1_PosValue; hw1.SlaveOperational := TRUE; hw2.RawPosIn := bench.Winch.COD2_PosValue; hw2.SlaveOperational := TRUE;
encoderM1(Enable := TRUE, HomingPermit := TRUE, HomingAtTargetM := btnM1, CfgHomingTargetM := 8.7, CfgTopSensorPosM := 8.7, HwIn := hw1, Cfg := cfgEncoder, Calib := calibM1); calibM1 := encoderM1.Calib;
bucketEdge(CLK := btnBucket);
encoderM2(Enable := TRUE, HomingPermit := TRUE, HomingAtTargetM := btnM2 OR bucketEdge.Q, CfgHomingTargetM := 23.7, CfgTopSensorPosM := 23.7, UseDynamicTarget := bucketEdge.Q, DynamicHomingTargetM := encoderM1.Measurement.CablePosM + cfgBucket.OffsetCloseM, HwIn := hw2, Cfg := cfgEncoder, Calib := calibM2); calibM2 := encoderM2.Calib;
bucket(Enable := TRUE, Mode := E_Mode.MAINT_N2, PowerContactorEngaged := TRUE, CablePosM1 := encoderM1.Measurement.CablePosM, CablePosM2 := encoderM2.Measurement.CablePosM, HomedM1 := encoderM1.Homed, HomedM2 := encoderM2.Homed, HomedAndReliableM1 := encoderM1.HomedAndReliable, HomedAndReliableM2 := encoderM2.HomedAndReliable, HomingSuspectM1 := encoderM1.HomingSuspect, HomingSuspectM2 := encoderM2.HomingSuspect, ConfirmClosePosition := btnBucket, Config := cfgBucket, BucketState := bucketState); bucketState := bucket.BucketState;
home.M1Status.HomedAndReliable := encoderM1.HomedAndReliable; home.M2Status.HomedAndReliable := encoderM2.HomedAndReliable; home(BucketOffsetValid := bucketState.BucketReferenced, BtnValidation := bench.Operator.JoyBtnRaw);
ADVANCE_TIME(10000000);
bench(M1_PresetTriggerCmd := encoderM1.HwOut.PresetTriggerCmd, M1_PresetValueOut := encoderM1.HwOut.PresetValueOut, M2_PresetTriggerCmd := encoderM2.HwOut.PresetTriggerCmd, M2_PresetValueOut := encoderM2.HwOut.PresetValueOut, RawPosM1 := raw1, RawPosM2 := raw2); raw1 := bench.RawPosM1; raw2 := bench.RawPosM2;
hw1.RawPosIn := bench.Winch.COD1_PosValue; hw1.SlaveOperational := TRUE; hw2.RawPosIn := bench.Winch.COD2_PosValue; hw2.SlaveOperational := TRUE;
encoderM1(Enable := TRUE, HomingPermit := TRUE, HomingAtTargetM := btnM1, CfgHomingTargetM := 8.7, CfgTopSensorPosM := 8.7, HwIn := hw1, Cfg := cfgEncoder, Calib := calibM1); calibM1 := encoderM1.Calib;
bucketEdge(CLK := btnBucket);
encoderM2(Enable := TRUE, HomingPermit := TRUE, HomingAtTargetM := btnM2 OR bucketEdge.Q, CfgHomingTargetM := 23.7, CfgTopSensorPosM := 23.7, UseDynamicTarget := bucketEdge.Q, DynamicHomingTargetM := encoderM1.Measurement.CablePosM + cfgBucket.OffsetCloseM, HwIn := hw2, Cfg := cfgEncoder, Calib := calibM2); calibM2 := encoderM2.Calib;
bucket(Enable := TRUE, Mode := E_Mode.MAINT_N2, PowerContactorEngaged := TRUE, CablePosM1 := encoderM1.Measurement.CablePosM, CablePosM2 := encoderM2.Measurement.CablePosM, HomedM1 := encoderM1.Homed, HomedM2 := encoderM2.Homed, HomedAndReliableM1 := encoderM1.HomedAndReliable, HomedAndReliableM2 := encoderM2.HomedAndReliable, HomingSuspectM1 := encoderM1.HomingSuspect, HomingSuspectM2 := encoderM2.HomingSuspect, ConfirmClosePosition := btnBucket, Config := cfgBucket, BucketState := bucketState); bucketState := bucket.BucketState;
home.M1Status.HomedAndReliable := encoderM1.HomedAndReliable; home.M2Status.HomedAndReliable := encoderM2.HomedAndReliable; home(BucketOffsetValid := bucketState.BucketReferenced, BtnValidation := bench.Operator.JoyBtnRaw);
ADVANCE_TIME(10000000);
bench(M1_PresetTriggerCmd := encoderM1.HwOut.PresetTriggerCmd, M1_PresetValueOut := encoderM1.HwOut.PresetValueOut, M2_PresetTriggerCmd := encoderM2.HwOut.PresetTriggerCmd, M2_PresetValueOut := encoderM2.HwOut.PresetValueOut, RawPosM1 := raw1, RawPosM2 := raw2); raw1 := bench.RawPosM1; raw2 := bench.RawPosM2;
hw1.RawPosIn := bench.Winch.COD1_PosValue; hw1.SlaveOperational := TRUE; hw2.RawPosIn := bench.Winch.COD2_PosValue; hw2.SlaveOperational := TRUE;
encoderM1(Enable := TRUE, HomingPermit := TRUE, HomingAtTargetM := btnM1, CfgHomingTargetM := 8.7, CfgTopSensorPosM := 8.7, HwIn := hw1, Cfg := cfgEncoder, Calib := calibM1); calibM1 := encoderM1.Calib;
bucketEdge(CLK := btnBucket);
encoderM2(Enable := TRUE, HomingPermit := TRUE, HomingAtTargetM := btnM2 OR bucketEdge.Q, CfgHomingTargetM := 23.7, CfgTopSensorPosM := 23.7, UseDynamicTarget := bucketEdge.Q, DynamicHomingTargetM := encoderM1.Measurement.CablePosM + cfgBucket.OffsetCloseM, HwIn := hw2, Cfg := cfgEncoder, Calib := calibM2); calibM2 := encoderM2.Calib;
bucket(Enable := TRUE, Mode := E_Mode.MAINT_N2, PowerContactorEngaged := TRUE, CablePosM1 := encoderM1.Measurement.CablePosM, CablePosM2 := encoderM2.Measurement.CablePosM, HomedM1 := encoderM1.Homed, HomedM2 := encoderM2.Homed, HomedAndReliableM1 := encoderM1.HomedAndReliable, HomedAndReliableM2 := encoderM2.HomedAndReliable, HomingSuspectM1 := encoderM1.HomingSuspect, HomingSuspectM2 := encoderM2.HomingSuspect, ConfirmClosePosition := btnBucket, Config := cfgBucket, BucketState := bucketState); bucketState := bucket.BucketState;
home.M1Status.HomedAndReliable := encoderM1.HomedAndReliable; home.M2Status.HomedAndReliable := encoderM2.HomedAndReliable; home(BucketOffsetValid := bucketState.BucketReferenced, BtnValidation := bench.Operator.JoyBtnRaw);
ADVANCE_TIME(10000000);
bench(M1_PresetTriggerCmd := encoderM1.HwOut.PresetTriggerCmd, M1_PresetValueOut := encoderM1.HwOut.PresetValueOut, M2_PresetTriggerCmd := encoderM2.HwOut.PresetTriggerCmd, M2_PresetValueOut := encoderM2.HwOut.PresetValueOut, RawPosM1 := raw1, RawPosM2 := raw2); raw1 := bench.RawPosM1; raw2 := bench.RawPosM2;
hw1.RawPosIn := bench.Winch.COD1_PosValue; hw1.SlaveOperational := TRUE; hw2.RawPosIn := bench.Winch.COD2_PosValue; hw2.SlaveOperational := TRUE;
encoderM1(Enable := TRUE, HomingPermit := TRUE, HomingAtTargetM := btnM1, CfgHomingTargetM := 8.7, CfgTopSensorPosM := 8.7, HwIn := hw1, Cfg := cfgEncoder, Calib := calibM1); calibM1 := encoderM1.Calib;
bucketEdge(CLK := btnBucket);
encoderM2(Enable := TRUE, HomingPermit := TRUE, HomingAtTargetM := btnM2 OR bucketEdge.Q, CfgHomingTargetM := 23.7, CfgTopSensorPosM := 23.7, UseDynamicTarget := bucketEdge.Q, DynamicHomingTargetM := encoderM1.Measurement.CablePosM + cfgBucket.OffsetCloseM, HwIn := hw2, Cfg := cfgEncoder, Calib := calibM2); calibM2 := encoderM2.Calib;
bucket(Enable := TRUE, Mode := E_Mode.MAINT_N2, PowerContactorEngaged := TRUE, CablePosM1 := encoderM1.Measurement.CablePosM, CablePosM2 := encoderM2.Measurement.CablePosM, HomedM1 := encoderM1.Homed, HomedM2 := encoderM2.Homed, HomedAndReliableM1 := encoderM1.HomedAndReliable, HomedAndReliableM2 := encoderM2.HomedAndReliable, HomingSuspectM1 := encoderM1.HomingSuspect, HomingSuspectM2 := encoderM2.HomingSuspect, ConfirmClosePosition := btnBucket, Config := cfgBucket, BucketState := bucketState); bucketState := bucket.BucketState;
home.M1Status.HomedAndReliable := encoderM1.HomedAndReliable; home.M2Status.HomedAndReliable := encoderM2.HomedAndReliable; home(BucketOffsetValid := bucketState.BucketReferenced, BtnValidation := bench.Operator.JoyBtnRaw);
ADVANCE_TIME(10000000);
bench(M1_PresetTriggerCmd := encoderM1.HwOut.PresetTriggerCmd, M1_PresetValueOut := encoderM1.HwOut.PresetValueOut, M2_PresetTriggerCmd := encoderM2.HwOut.PresetTriggerCmd, M2_PresetValueOut := encoderM2.HwOut.PresetValueOut, RawPosM1 := raw1, RawPosM2 := raw2); raw1 := bench.RawPosM1; raw2 := bench.RawPosM2;
hw1.RawPosIn := bench.Winch.COD1_PosValue; hw1.SlaveOperational := TRUE; hw2.RawPosIn := bench.Winch.COD2_PosValue; hw2.SlaveOperational := TRUE;
encoderM1(Enable := TRUE, HomingPermit := TRUE, HomingAtTargetM := btnM1, CfgHomingTargetM := 8.7, CfgTopSensorPosM := 8.7, HwIn := hw1, Cfg := cfgEncoder, Calib := calibM1); calibM1 := encoderM1.Calib;
bucketEdge(CLK := btnBucket);
encoderM2(Enable := TRUE, HomingPermit := TRUE, HomingAtTargetM := btnM2 OR bucketEdge.Q, CfgHomingTargetM := 23.7, CfgTopSensorPosM := 23.7, UseDynamicTarget := bucketEdge.Q, DynamicHomingTargetM := encoderM1.Measurement.CablePosM + cfgBucket.OffsetCloseM, HwIn := hw2, Cfg := cfgEncoder, Calib := calibM2); calibM2 := encoderM2.Calib;
bucket(Enable := TRUE, Mode := E_Mode.MAINT_N2, PowerContactorEngaged := TRUE, CablePosM1 := encoderM1.Measurement.CablePosM, CablePosM2 := encoderM2.Measurement.CablePosM, HomedM1 := encoderM1.Homed, HomedM2 := encoderM2.Homed, HomedAndReliableM1 := encoderM1.HomedAndReliable, HomedAndReliableM2 := encoderM2.HomedAndReliable, HomingSuspectM1 := encoderM1.HomingSuspect, HomingSuspectM2 := encoderM2.HomingSuspect, ConfirmClosePosition := btnBucket, Config := cfgBucket, BucketState := bucketState); bucketState := bucket.BucketState;
home.M1Status.HomedAndReliable := encoderM1.HomedAndReliable; home.M2Status.HomedAndReliable := encoderM2.HomedAndReliable; home(BucketOffsetValid := bucketState.BucketReferenced, BtnValidation := bench.Operator.JoyBtnRaw);
ADVANCE_TIME(10000000);
bench(M1_PresetTriggerCmd := encoderM1.HwOut.PresetTriggerCmd, M1_PresetValueOut := encoderM1.HwOut.PresetValueOut, M2_PresetTriggerCmd := encoderM2.HwOut.PresetTriggerCmd, M2_PresetValueOut := encoderM2.HwOut.PresetValueOut, RawPosM1 := raw1, RawPosM2 := raw2); raw1 := bench.RawPosM1; raw2 := bench.RawPosM2;
hw1.RawPosIn := bench.Winch.COD1_PosValue; hw1.SlaveOperational := TRUE; hw2.RawPosIn := bench.Winch.COD2_PosValue; hw2.SlaveOperational := TRUE;
encoderM1(Enable := TRUE, HomingPermit := TRUE, HomingAtTargetM := btnM1, CfgHomingTargetM := 8.7, CfgTopSensorPosM := 8.7, HwIn := hw1, Cfg := cfgEncoder, Calib := calibM1); calibM1 := encoderM1.Calib;
bucketEdge(CLK := btnBucket);
encoderM2(Enable := TRUE, HomingPermit := TRUE, HomingAtTargetM := btnM2 OR bucketEdge.Q, CfgHomingTargetM := 23.7, CfgTopSensorPosM := 23.7, UseDynamicTarget := bucketEdge.Q, DynamicHomingTargetM := encoderM1.Measurement.CablePosM + cfgBucket.OffsetCloseM, HwIn := hw2, Cfg := cfgEncoder, Calib := calibM2); calibM2 := encoderM2.Calib;
bucket(Enable := TRUE, Mode := E_Mode.MAINT_N2, PowerContactorEngaged := TRUE, CablePosM1 := encoderM1.Measurement.CablePosM, CablePosM2 := encoderM2.Measurement.CablePosM, HomedM1 := encoderM1.Homed, HomedM2 := encoderM2.Homed, HomedAndReliableM1 := encoderM1.HomedAndReliable, HomedAndReliableM2 := encoderM2.HomedAndReliable, HomingSuspectM1 := encoderM1.HomingSuspect, HomingSuspectM2 := encoderM2.HomingSuspect, ConfirmClosePosition := btnBucket, Config := cfgBucket, BucketState := bucketState); bucketState := bucket.BucketState;
home.M1Status.HomedAndReliable := encoderM1.HomedAndReliable; home.M2Status.HomedAndReliable := encoderM2.HomedAndReliable; home(BucketOffsetValid := bucketState.BucketReferenced, BtnValidation := bench.Operator.JoyBtnRaw);
ADVANCE_TIME(10000000);
bench(M1_PresetTriggerCmd := encoderM1.HwOut.PresetTriggerCmd, M1_PresetValueOut := encoderM1.HwOut.PresetValueOut, M2_PresetTriggerCmd := encoderM2.HwOut.PresetTriggerCmd, M2_PresetValueOut := encoderM2.HwOut.PresetValueOut, RawPosM1 := raw1, RawPosM2 := raw2); raw1 := bench.RawPosM1; raw2 := bench.RawPosM2;
hw1.RawPosIn := bench.Winch.COD1_PosValue; hw1.SlaveOperational := TRUE; hw2.RawPosIn := bench.Winch.COD2_PosValue; hw2.SlaveOperational := TRUE;
encoderM1(Enable := TRUE, HomingPermit := TRUE, HomingAtTargetM := btnM1, CfgHomingTargetM := 8.7, CfgTopSensorPosM := 8.7, HwIn := hw1, Cfg := cfgEncoder, Calib := calibM1); calibM1 := encoderM1.Calib;
bucketEdge(CLK := btnBucket);
encoderM2(Enable := TRUE, HomingPermit := TRUE, HomingAtTargetM := btnM2 OR bucketEdge.Q, CfgHomingTargetM := 23.7, CfgTopSensorPosM := 23.7, UseDynamicTarget := bucketEdge.Q, DynamicHomingTargetM := encoderM1.Measurement.CablePosM + cfgBucket.OffsetCloseM, HwIn := hw2, Cfg := cfgEncoder, Calib := calibM2); calibM2 := encoderM2.Calib;
bucket(Enable := TRUE, Mode := E_Mode.MAINT_N2, PowerContactorEngaged := TRUE, CablePosM1 := encoderM1.Measurement.CablePosM, CablePosM2 := encoderM2.Measurement.CablePosM, HomedM1 := encoderM1.Homed, HomedM2 := encoderM2.Homed, HomedAndReliableM1 := encoderM1.HomedAndReliable, HomedAndReliableM2 := encoderM2.HomedAndReliable, HomingSuspectM1 := encoderM1.HomingSuspect, HomingSuspectM2 := encoderM2.HomingSuspect, ConfirmClosePosition := btnBucket, Config := cfgBucket, BucketState := bucketState); bucketState := bucket.BucketState;
home.M1Status.HomedAndReliable := encoderM1.HomedAndReliable; home.M2Status.HomedAndReliable := encoderM2.HomedAndReliable; home(BucketOffsetValid := bucketState.BucketReferenced, BtnValidation := bench.Operator.JoyBtnRaw);
ADVANCE_TIME(10000000);
bench(M1_PresetTriggerCmd := encoderM1.HwOut.PresetTriggerCmd, M1_PresetValueOut := encoderM1.HwOut.PresetValueOut, M2_PresetTriggerCmd := encoderM2.HwOut.PresetTriggerCmd, M2_PresetValueOut := encoderM2.HwOut.PresetValueOut, RawPosM1 := raw1, RawPosM2 := raw2); raw1 := bench.RawPosM1; raw2 := bench.RawPosM2;
hw1.RawPosIn := bench.Winch.COD1_PosValue; hw1.SlaveOperational := TRUE; hw2.RawPosIn := bench.Winch.COD2_PosValue; hw2.SlaveOperational := TRUE;
encoderM1(Enable := TRUE, HomingPermit := TRUE, HomingAtTargetM := btnM1, CfgHomingTargetM := 8.7, CfgTopSensorPosM := 8.7, HwIn := hw1, Cfg := cfgEncoder, Calib := calibM1); calibM1 := encoderM1.Calib;
bucketEdge(CLK := btnBucket);
encoderM2(Enable := TRUE, HomingPermit := TRUE, HomingAtTargetM := btnM2 OR bucketEdge.Q, CfgHomingTargetM := 23.7, CfgTopSensorPosM := 23.7, UseDynamicTarget := bucketEdge.Q, DynamicHomingTargetM := encoderM1.Measurement.CablePosM + cfgBucket.OffsetCloseM, HwIn := hw2, Cfg := cfgEncoder, Calib := calibM2); calibM2 := encoderM2.Calib;
bucket(Enable := TRUE, Mode := E_Mode.MAINT_N2, PowerContactorEngaged := TRUE, CablePosM1 := encoderM1.Measurement.CablePosM, CablePosM2 := encoderM2.Measurement.CablePosM, HomedM1 := encoderM1.Homed, HomedM2 := encoderM2.Homed, HomedAndReliableM1 := encoderM1.HomedAndReliable, HomedAndReliableM2 := encoderM2.HomedAndReliable, HomingSuspectM1 := encoderM1.HomingSuspect, HomingSuspectM2 := encoderM2.HomingSuspect, ConfirmClosePosition := btnBucket, Config := cfgBucket, BucketState := bucketState); bucketState := bucket.BucketState;
home.M1Status.HomedAndReliable := encoderM1.HomedAndReliable; home.M2Status.HomedAndReliable := encoderM2.HomedAndReliable; home(BucketOffsetValid := bucketState.BucketReferenced, BtnValidation := bench.Operator.JoyBtnRaw);
ADVANCE_TIME(10000000);
bench(M1_PresetTriggerCmd := encoderM1.HwOut.PresetTriggerCmd, M1_PresetValueOut := encoderM1.HwOut.PresetValueOut, M2_PresetTriggerCmd := encoderM2.HwOut.PresetTriggerCmd, M2_PresetValueOut := encoderM2.HwOut.PresetValueOut, RawPosM1 := raw1, RawPosM2 := raw2); raw1 := bench.RawPosM1; raw2 := bench.RawPosM2;
hw1.RawPosIn := bench.Winch.COD1_PosValue; hw1.SlaveOperational := TRUE; hw2.RawPosIn := bench.Winch.COD2_PosValue; hw2.SlaveOperational := TRUE;
encoderM1(Enable := TRUE, HomingPermit := TRUE, HomingAtTargetM := btnM1, CfgHomingTargetM := 8.7, CfgTopSensorPosM := 8.7, HwIn := hw1, Cfg := cfgEncoder, Calib := calibM1); calibM1 := encoderM1.Calib;
bucketEdge(CLK := btnBucket);
encoderM2(Enable := TRUE, HomingPermit := TRUE, HomingAtTargetM := btnM2 OR bucketEdge.Q, CfgHomingTargetM := 23.7, CfgTopSensorPosM := 23.7, UseDynamicTarget := bucketEdge.Q, DynamicHomingTargetM := encoderM1.Measurement.CablePosM + cfgBucket.OffsetCloseM, HwIn := hw2, Cfg := cfgEncoder, Calib := calibM2); calibM2 := encoderM2.Calib;
bucket(Enable := TRUE, Mode := E_Mode.MAINT_N2, PowerContactorEngaged := TRUE, CablePosM1 := encoderM1.Measurement.CablePosM, CablePosM2 := encoderM2.Measurement.CablePosM, HomedM1 := encoderM1.Homed, HomedM2 := encoderM2.Homed, HomedAndReliableM1 := encoderM1.HomedAndReliable, HomedAndReliableM2 := encoderM2.HomedAndReliable, HomingSuspectM1 := encoderM1.HomingSuspect, HomingSuspectM2 := encoderM2.HomingSuspect, ConfirmClosePosition := btnBucket, Config := cfgBucket, BucketState := bucketState); bucketState := bucket.BucketState;
home.M1Status.HomedAndReliable := encoderM1.HomedAndReliable; home.M2Status.HomedAndReliable := encoderM2.HomedAndReliable; home(BucketOffsetValid := bucketState.BucketReferenced, BtnValidation := bench.Operator.JoyBtnRaw);
ADVANCE_TIME(10000000);
bench(M1_PresetTriggerCmd := encoderM1.HwOut.PresetTriggerCmd, M1_PresetValueOut := encoderM1.HwOut.PresetValueOut, M2_PresetTriggerCmd := encoderM2.HwOut.PresetTriggerCmd, M2_PresetValueOut := encoderM2.HwOut.PresetValueOut, RawPosM1 := raw1, RawPosM2 := raw2); raw1 := bench.RawPosM1; raw2 := bench.RawPosM2;
hw1.RawPosIn := bench.Winch.COD1_PosValue; hw1.SlaveOperational := TRUE; hw2.RawPosIn := bench.Winch.COD2_PosValue; hw2.SlaveOperational := TRUE;
encoderM1(Enable := TRUE, HomingPermit := TRUE, HomingAtTargetM := btnM1, CfgHomingTargetM := 8.7, CfgTopSensorPosM := 8.7, HwIn := hw1, Cfg := cfgEncoder, Calib := calibM1); calibM1 := encoderM1.Calib;
bucketEdge(CLK := btnBucket);
encoderM2(Enable := TRUE, HomingPermit := TRUE, HomingAtTargetM := btnM2 OR bucketEdge.Q, CfgHomingTargetM := 23.7, CfgTopSensorPosM := 23.7, UseDynamicTarget := bucketEdge.Q, DynamicHomingTargetM := encoderM1.Measurement.CablePosM + cfgBucket.OffsetCloseM, HwIn := hw2, Cfg := cfgEncoder, Calib := calibM2); calibM2 := encoderM2.Calib;
bucket(Enable := TRUE, Mode := E_Mode.MAINT_N2, PowerContactorEngaged := TRUE, CablePosM1 := encoderM1.Measurement.CablePosM, CablePosM2 := encoderM2.Measurement.CablePosM, HomedM1 := encoderM1.Homed, HomedM2 := encoderM2.Homed, HomedAndReliableM1 := encoderM1.HomedAndReliable, HomedAndReliableM2 := encoderM2.HomedAndReliable, HomingSuspectM1 := encoderM1.HomingSuspect, HomingSuspectM2 := encoderM2.HomingSuspect, ConfirmClosePosition := btnBucket, Config := cfgBucket, BucketState := bucketState); bucketState := bucket.BucketState;
home.M1Status.HomedAndReliable := encoderM1.HomedAndReliable; home.M2Status.HomedAndReliable := encoderM2.HomedAndReliable; home(BucketOffsetValid := bucketState.BucketReferenced, BtnValidation := bench.Operator.JoyBtnRaw);
ADVANCE_TIME(10000000);
bench(M1_PresetTriggerCmd := encoderM1.HwOut.PresetTriggerCmd, M1_PresetValueOut := encoderM1.HwOut.PresetValueOut, M2_PresetTriggerCmd := encoderM2.HwOut.PresetTriggerCmd, M2_PresetValueOut := encoderM2.HwOut.PresetValueOut, RawPosM1 := raw1, RawPosM2 := raw2); raw1 := bench.RawPosM1; raw2 := bench.RawPosM2;
hw1.RawPosIn := bench.Winch.COD1_PosValue; hw1.SlaveOperational := TRUE; hw2.RawPosIn := bench.Winch.COD2_PosValue; hw2.SlaveOperational := TRUE;
encoderM1(Enable := TRUE, HomingPermit := TRUE, HomingAtTargetM := btnM1, CfgHomingTargetM := 8.7, CfgTopSensorPosM := 8.7, HwIn := hw1, Cfg := cfgEncoder, Calib := calibM1); calibM1 := encoderM1.Calib;
bucketEdge(CLK := btnBucket);
encoderM2(Enable := TRUE, HomingPermit := TRUE, HomingAtTargetM := btnM2 OR bucketEdge.Q, CfgHomingTargetM := 23.7, CfgTopSensorPosM := 23.7, UseDynamicTarget := bucketEdge.Q, DynamicHomingTargetM := encoderM1.Measurement.CablePosM + cfgBucket.OffsetCloseM, HwIn := hw2, Cfg := cfgEncoder, Calib := calibM2); calibM2 := encoderM2.Calib;
bucket(Enable := TRUE, Mode := E_Mode.MAINT_N2, PowerContactorEngaged := TRUE, CablePosM1 := encoderM1.Measurement.CablePosM, CablePosM2 := encoderM2.Measurement.CablePosM, HomedM1 := encoderM1.Homed, HomedM2 := encoderM2.Homed, HomedAndReliableM1 := encoderM1.HomedAndReliable, HomedAndReliableM2 := encoderM2.HomedAndReliable, HomingSuspectM1 := encoderM1.HomingSuspect, HomingSuspectM2 := encoderM2.HomingSuspect, ConfirmClosePosition := btnBucket, Config := cfgBucket, BucketState := bucketState); bucketState := bucket.BucketState;
home.M1Status.HomedAndReliable := encoderM1.HomedAndReliable; home.M2Status.HomedAndReliable := encoderM2.HomedAndReliable; home(BucketOffsetValid := bucketState.BucketReferenced, BtnValidation := bench.Operator.JoyBtnRaw);
ADVANCE_TIME(10000000);
bench(M1_PresetTriggerCmd := encoderM1.HwOut.PresetTriggerCmd, M1_PresetValueOut := encoderM1.HwOut.PresetValueOut, M2_PresetTriggerCmd := encoderM2.HwOut.PresetTriggerCmd, M2_PresetValueOut := encoderM2.HwOut.PresetValueOut, RawPosM1 := raw1, RawPosM2 := raw2); raw1 := bench.RawPosM1; raw2 := bench.RawPosM2;
hw1.RawPosIn := bench.Winch.COD1_PosValue; hw1.SlaveOperational := TRUE; hw2.RawPosIn := bench.Winch.COD2_PosValue; hw2.SlaveOperational := TRUE;
encoderM1(Enable := TRUE, HomingPermit := TRUE, HomingAtTargetM := btnM1, CfgHomingTargetM := 8.7, CfgTopSensorPosM := 8.7, HwIn := hw1, Cfg := cfgEncoder, Calib := calibM1); calibM1 := encoderM1.Calib;
bucketEdge(CLK := btnBucket);
encoderM2(Enable := TRUE, HomingPermit := TRUE, HomingAtTargetM := btnM2 OR bucketEdge.Q, CfgHomingTargetM := 23.7, CfgTopSensorPosM := 23.7, UseDynamicTarget := bucketEdge.Q, DynamicHomingTargetM := encoderM1.Measurement.CablePosM + cfgBucket.OffsetCloseM, HwIn := hw2, Cfg := cfgEncoder, Calib := calibM2); calibM2 := encoderM2.Calib;
bucket(Enable := TRUE, Mode := E_Mode.MAINT_N2, PowerContactorEngaged := TRUE, CablePosM1 := encoderM1.Measurement.CablePosM, CablePosM2 := encoderM2.Measurement.CablePosM, HomedM1 := encoderM1.Homed, HomedM2 := encoderM2.Homed, HomedAndReliableM1 := encoderM1.HomedAndReliable, HomedAndReliableM2 := encoderM2.HomedAndReliable, HomingSuspectM1 := encoderM1.HomingSuspect, HomingSuspectM2 := encoderM2.HomingSuspect, ConfirmClosePosition := btnBucket, Config := cfgBucket, BucketState := bucketState); bucketState := bucket.BucketState;
home.M1Status.HomedAndReliable := encoderM1.HomedAndReliable; home.M2Status.HomedAndReliable := encoderM2.HomedAndReliable; home(BucketOffsetValid := bucketState.BucketReferenced, BtnValidation := bench.Operator.JoyBtnRaw);
ADVANCE_TIME(10000000);
bench(M1_PresetTriggerCmd := encoderM1.HwOut.PresetTriggerCmd, M1_PresetValueOut := encoderM1.HwOut.PresetValueOut, M2_PresetTriggerCmd := encoderM2.HwOut.PresetTriggerCmd, M2_PresetValueOut := encoderM2.HwOut.PresetValueOut, RawPosM1 := raw1, RawPosM2 := raw2); raw1 := bench.RawPosM1; raw2 := bench.RawPosM2;
hw1.RawPosIn := bench.Winch.COD1_PosValue; hw1.SlaveOperational := TRUE; hw2.RawPosIn := bench.Winch.COD2_PosValue; hw2.SlaveOperational := TRUE;
encoderM1(Enable := TRUE, HomingPermit := TRUE, HomingAtTargetM := btnM1, CfgHomingTargetM := 8.7, CfgTopSensorPosM := 8.7, HwIn := hw1, Cfg := cfgEncoder, Calib := calibM1); calibM1 := encoderM1.Calib;
bucketEdge(CLK := btnBucket);
encoderM2(Enable := TRUE, HomingPermit := TRUE, HomingAtTargetM := btnM2 OR bucketEdge.Q, CfgHomingTargetM := 23.7, CfgTopSensorPosM := 23.7, UseDynamicTarget := bucketEdge.Q, DynamicHomingTargetM := encoderM1.Measurement.CablePosM + cfgBucket.OffsetCloseM, HwIn := hw2, Cfg := cfgEncoder, Calib := calibM2); calibM2 := encoderM2.Calib;
bucket(Enable := TRUE, Mode := E_Mode.MAINT_N2, PowerContactorEngaged := TRUE, CablePosM1 := encoderM1.Measurement.CablePosM, CablePosM2 := encoderM2.Measurement.CablePosM, HomedM1 := encoderM1.Homed, HomedM2 := encoderM2.Homed, HomedAndReliableM1 := encoderM1.HomedAndReliable, HomedAndReliableM2 := encoderM2.HomedAndReliable, HomingSuspectM1 := encoderM1.HomingSuspect, HomingSuspectM2 := encoderM2.HomingSuspect, ConfirmClosePosition := btnBucket, Config := cfgBucket, BucketState := bucketState); bucketState := bucket.BucketState;
home.M1Status.HomedAndReliable := encoderM1.HomedAndReliable; home.M2Status.HomedAndReliable := encoderM2.HomedAndReliable; home(BucketOffsetValid := bucketState.BucketReferenced, BtnValidation := bench.Operator.JoyBtnRaw);
ADVANCE_TIME(10000000);
bench(M1_PresetTriggerCmd := encoderM1.HwOut.PresetTriggerCmd, M1_PresetValueOut := encoderM1.HwOut.PresetValueOut, M2_PresetTriggerCmd := encoderM2.HwOut.PresetTriggerCmd, M2_PresetValueOut := encoderM2.HwOut.PresetValueOut, RawPosM1 := raw1, RawPosM2 := raw2); raw1 := bench.RawPosM1; raw2 := bench.RawPosM2;
hw1.RawPosIn := bench.Winch.COD1_PosValue; hw1.SlaveOperational := TRUE; hw2.RawPosIn := bench.Winch.COD2_PosValue; hw2.SlaveOperational := TRUE;
encoderM1(Enable := TRUE, HomingPermit := TRUE, HomingAtTargetM := btnM1, CfgHomingTargetM := 8.7, CfgTopSensorPosM := 8.7, HwIn := hw1, Cfg := cfgEncoder, Calib := calibM1); calibM1 := encoderM1.Calib;
bucketEdge(CLK := btnBucket);
encoderM2(Enable := TRUE, HomingPermit := TRUE, HomingAtTargetM := btnM2 OR bucketEdge.Q, CfgHomingTargetM := 23.7, CfgTopSensorPosM := 23.7, UseDynamicTarget := bucketEdge.Q, DynamicHomingTargetM := encoderM1.Measurement.CablePosM + cfgBucket.OffsetCloseM, HwIn := hw2, Cfg := cfgEncoder, Calib := calibM2); calibM2 := encoderM2.Calib;
bucket(Enable := TRUE, Mode := E_Mode.MAINT_N2, PowerContactorEngaged := TRUE, CablePosM1 := encoderM1.Measurement.CablePosM, CablePosM2 := encoderM2.Measurement.CablePosM, HomedM1 := encoderM1.Homed, HomedM2 := encoderM2.Homed, HomedAndReliableM1 := encoderM1.HomedAndReliable, HomedAndReliableM2 := encoderM2.HomedAndReliable, HomingSuspectM1 := encoderM1.HomingSuspect, HomingSuspectM2 := encoderM2.HomingSuspect, ConfirmClosePosition := btnBucket, Config := cfgBucket, BucketState := bucketState); bucketState := bucket.BucketState;
home.M1Status.HomedAndReliable := encoderM1.HomedAndReliable; home.M2Status.HomedAndReliable := encoderM2.HomedAndReliable; home(BucketOffsetValid := bucketState.BucketReferenced, BtnValidation := bench.Operator.JoyBtnRaw);
ADVANCE_TIME(10000000);
bench(M1_PresetTriggerCmd := encoderM1.HwOut.PresetTriggerCmd, M1_PresetValueOut := encoderM1.HwOut.PresetValueOut, M2_PresetTriggerCmd := encoderM2.HwOut.PresetTriggerCmd, M2_PresetValueOut := encoderM2.HwOut.PresetValueOut, RawPosM1 := raw1, RawPosM2 := raw2); raw1 := bench.RawPosM1; raw2 := bench.RawPosM2;
hw1.RawPosIn := bench.Winch.COD1_PosValue; hw1.SlaveOperational := TRUE; hw2.RawPosIn := bench.Winch.COD2_PosValue; hw2.SlaveOperational := TRUE;
encoderM1(Enable := TRUE, HomingPermit := TRUE, HomingAtTargetM := btnM1, CfgHomingTargetM := 8.7, CfgTopSensorPosM := 8.7, HwIn := hw1, Cfg := cfgEncoder, Calib := calibM1); calibM1 := encoderM1.Calib;
bucketEdge(CLK := btnBucket);
encoderM2(Enable := TRUE, HomingPermit := TRUE, HomingAtTargetM := btnM2 OR bucketEdge.Q, CfgHomingTargetM := 23.7, CfgTopSensorPosM := 23.7, UseDynamicTarget := bucketEdge.Q, DynamicHomingTargetM := encoderM1.Measurement.CablePosM + cfgBucket.OffsetCloseM, HwIn := hw2, Cfg := cfgEncoder, Calib := calibM2); calibM2 := encoderM2.Calib;
bucket(Enable := TRUE, Mode := E_Mode.MAINT_N2, PowerContactorEngaged := TRUE, CablePosM1 := encoderM1.Measurement.CablePosM, CablePosM2 := encoderM2.Measurement.CablePosM, HomedM1 := encoderM1.Homed, HomedM2 := encoderM2.Homed, HomedAndReliableM1 := encoderM1.HomedAndReliable, HomedAndReliableM2 := encoderM2.HomedAndReliable, HomingSuspectM1 := encoderM1.HomingSuspect, HomingSuspectM2 := encoderM2.HomingSuspect, ConfirmClosePosition := btnBucket, Config := cfgBucket, BucketState := bucketState); bucketState := bucket.BucketState;
home.M1Status.HomedAndReliable := encoderM1.HomedAndReliable; home.M2Status.HomedAndReliable := encoderM2.HomedAndReliable; home(BucketOffsetValid := bucketState.BucketReferenced, BtnValidation := bench.Operator.JoyBtnRaw);
ADVANCE_TIME(10000000);
bench(M1_PresetTriggerCmd := encoderM1.HwOut.PresetTriggerCmd, M1_PresetValueOut := encoderM1.HwOut.PresetValueOut, M2_PresetTriggerCmd := encoderM2.HwOut.PresetTriggerCmd, M2_PresetValueOut := encoderM2.HwOut.PresetValueOut, RawPosM1 := raw1, RawPosM2 := raw2); raw1 := bench.RawPosM1; raw2 := bench.RawPosM2;
hw1.RawPosIn := bench.Winch.COD1_PosValue; hw1.SlaveOperational := TRUE; hw2.RawPosIn := bench.Winch.COD2_PosValue; hw2.SlaveOperational := TRUE;
encoderM1(Enable := TRUE, HomingPermit := TRUE, HomingAtTargetM := btnM1, CfgHomingTargetM := 8.7, CfgTopSensorPosM := 8.7, HwIn := hw1, Cfg := cfgEncoder, Calib := calibM1); calibM1 := encoderM1.Calib;
bucketEdge(CLK := btnBucket);
encoderM2(Enable := TRUE, HomingPermit := TRUE, HomingAtTargetM := btnM2 OR bucketEdge.Q, CfgHomingTargetM := 23.7, CfgTopSensorPosM := 23.7, UseDynamicTarget := bucketEdge.Q, DynamicHomingTargetM := encoderM1.Measurement.CablePosM + cfgBucket.OffsetCloseM, HwIn := hw2, Cfg := cfgEncoder, Calib := calibM2); calibM2 := encoderM2.Calib;
bucket(Enable := TRUE, Mode := E_Mode.MAINT_N2, PowerContactorEngaged := TRUE, CablePosM1 := encoderM1.Measurement.CablePosM, CablePosM2 := encoderM2.Measurement.CablePosM, HomedM1 := encoderM1.Homed, HomedM2 := encoderM2.Homed, HomedAndReliableM1 := encoderM1.HomedAndReliable, HomedAndReliableM2 := encoderM2.HomedAndReliable, HomingSuspectM1 := encoderM1.HomingSuspect, HomingSuspectM2 := encoderM2.HomingSuspect, ConfirmClosePosition := btnBucket, Config := cfgBucket, BucketState := bucketState); bucketState := bucket.BucketState;
home.M1Status.HomedAndReliable := encoderM1.HomedAndReliable; home.M2Status.HomedAndReliable := encoderM2.HomedAndReliable; home(BucketOffsetValid := bucketState.BucketReferenced, BtnValidation := bench.Operator.JoyBtnRaw);
ADVANCE_TIME(10000000);
bench(M1_PresetTriggerCmd := encoderM1.HwOut.PresetTriggerCmd, M1_PresetValueOut := encoderM1.HwOut.PresetValueOut, M2_PresetTriggerCmd := encoderM2.HwOut.PresetTriggerCmd, M2_PresetValueOut := encoderM2.HwOut.PresetValueOut, RawPosM1 := raw1, RawPosM2 := raw2); raw1 := bench.RawPosM1; raw2 := bench.RawPosM2;
hw1.RawPosIn := bench.Winch.COD1_PosValue; hw1.SlaveOperational := TRUE; hw2.RawPosIn := bench.Winch.COD2_PosValue; hw2.SlaveOperational := TRUE;
encoderM1(Enable := TRUE, HomingPermit := TRUE, HomingAtTargetM := btnM1, CfgHomingTargetM := 8.7, CfgTopSensorPosM := 8.7, HwIn := hw1, Cfg := cfgEncoder, Calib := calibM1); calibM1 := encoderM1.Calib;
bucketEdge(CLK := btnBucket);
encoderM2(Enable := TRUE, HomingPermit := TRUE, HomingAtTargetM := btnM2 OR bucketEdge.Q, CfgHomingTargetM := 23.7, CfgTopSensorPosM := 23.7, UseDynamicTarget := bucketEdge.Q, DynamicHomingTargetM := encoderM1.Measurement.CablePosM + cfgBucket.OffsetCloseM, HwIn := hw2, Cfg := cfgEncoder, Calib := calibM2); calibM2 := encoderM2.Calib;
bucket(Enable := TRUE, Mode := E_Mode.MAINT_N2, PowerContactorEngaged := TRUE, CablePosM1 := encoderM1.Measurement.CablePosM, CablePosM2 := encoderM2.Measurement.CablePosM, HomedM1 := encoderM1.Homed, HomedM2 := encoderM2.Homed, HomedAndReliableM1 := encoderM1.HomedAndReliable, HomedAndReliableM2 := encoderM2.HomedAndReliable, HomingSuspectM1 := encoderM1.HomingSuspect, HomingSuspectM2 := encoderM2.HomingSuspect, ConfirmClosePosition := btnBucket, Config := cfgBucket, BucketState := bucketState); bucketState := bucket.BucketState;
home.M1Status.HomedAndReliable := encoderM1.HomedAndReliable; home.M2Status.HomedAndReliable := encoderM2.HomedAndReliable; home(BucketOffsetValid := bucketState.BucketReferenced, BtnValidation := bench.Operator.JoyBtnRaw);
ADVANCE_TIME(10000000);
bench(M1_PresetTriggerCmd := encoderM1.HwOut.PresetTriggerCmd, M1_PresetValueOut := encoderM1.HwOut.PresetValueOut, M2_PresetTriggerCmd := encoderM2.HwOut.PresetTriggerCmd, M2_PresetValueOut := encoderM2.HwOut.PresetValueOut, RawPosM1 := raw1, RawPosM2 := raw2); raw1 := bench.RawPosM1; raw2 := bench.RawPosM2;
hw1.RawPosIn := bench.Winch.COD1_PosValue; hw1.SlaveOperational := TRUE; hw2.RawPosIn := bench.Winch.COD2_PosValue; hw2.SlaveOperational := TRUE;
encoderM1(Enable := TRUE, HomingPermit := TRUE, HomingAtTargetM := btnM1, CfgHomingTargetM := 8.7, CfgTopSensorPosM := 8.7, HwIn := hw1, Cfg := cfgEncoder, Calib := calibM1); calibM1 := encoderM1.Calib;
bucketEdge(CLK := btnBucket);
encoderM2(Enable := TRUE, HomingPermit := TRUE, HomingAtTargetM := btnM2 OR bucketEdge.Q, CfgHomingTargetM := 23.7, CfgTopSensorPosM := 23.7, UseDynamicTarget := bucketEdge.Q, DynamicHomingTargetM := encoderM1.Measurement.CablePosM + cfgBucket.OffsetCloseM, HwIn := hw2, Cfg := cfgEncoder, Calib := calibM2); calibM2 := encoderM2.Calib;
bucket(Enable := TRUE, Mode := E_Mode.MAINT_N2, PowerContactorEngaged := TRUE, CablePosM1 := encoderM1.Measurement.CablePosM, CablePosM2 := encoderM2.Measurement.CablePosM, HomedM1 := encoderM1.Homed, HomedM2 := encoderM2.Homed, HomedAndReliableM1 := encoderM1.HomedAndReliable, HomedAndReliableM2 := encoderM2.HomedAndReliable, HomingSuspectM1 := encoderM1.HomingSuspect, HomingSuspectM2 := encoderM2.HomingSuspect, ConfirmClosePosition := btnBucket, Config := cfgBucket, BucketState := bucketState); bucketState := bucket.BucketState;
home.M1Status.HomedAndReliable := encoderM1.HomedAndReliable; home.M2Status.HomedAndReliable := encoderM2.HomedAndReliable; home(BucketOffsetValid := bucketState.BucketReferenced, BtnValidation := bench.Operator.JoyBtnRaw);
ADVANCE_TIME(10000000);
bench(M1_PresetTriggerCmd := encoderM1.HwOut.PresetTriggerCmd, M1_PresetValueOut := encoderM1.HwOut.PresetValueOut, M2_PresetTriggerCmd := encoderM2.HwOut.PresetTriggerCmd, M2_PresetValueOut := encoderM2.HwOut.PresetValueOut, RawPosM1 := raw1, RawPosM2 := raw2); raw1 := bench.RawPosM1; raw2 := bench.RawPosM2;
hw1.RawPosIn := bench.Winch.COD1_PosValue; hw1.SlaveOperational := TRUE; hw2.RawPosIn := bench.Winch.COD2_PosValue; hw2.SlaveOperational := TRUE;
encoderM1(Enable := TRUE, HomingPermit := TRUE, HomingAtTargetM := btnM1, CfgHomingTargetM := 8.7, CfgTopSensorPosM := 8.7, HwIn := hw1, Cfg := cfgEncoder, Calib := calibM1); calibM1 := encoderM1.Calib;
bucketEdge(CLK := btnBucket);
encoderM2(Enable := TRUE, HomingPermit := TRUE, HomingAtTargetM := btnM2 OR bucketEdge.Q, CfgHomingTargetM := 23.7, CfgTopSensorPosM := 23.7, UseDynamicTarget := bucketEdge.Q, DynamicHomingTargetM := encoderM1.Measurement.CablePosM + cfgBucket.OffsetCloseM, HwIn := hw2, Cfg := cfgEncoder, Calib := calibM2); calibM2 := encoderM2.Calib;
bucket(Enable := TRUE, Mode := E_Mode.MAINT_N2, PowerContactorEngaged := TRUE, CablePosM1 := encoderM1.Measurement.CablePosM, CablePosM2 := encoderM2.Measurement.CablePosM, HomedM1 := encoderM1.Homed, HomedM2 := encoderM2.Homed, HomedAndReliableM1 := encoderM1.HomedAndReliable, HomedAndReliableM2 := encoderM2.HomedAndReliable, HomingSuspectM1 := encoderM1.HomingSuspect, HomingSuspectM2 := encoderM2.HomingSuspect, ConfirmClosePosition := btnBucket, Config := cfgBucket, BucketState := bucketState); bucketState := bucket.BucketState;
home.M1Status.HomedAndReliable := encoderM1.HomedAndReliable; home.M2Status.HomedAndReliable := encoderM2.HomedAndReliable; home(BucketOffsetValid := bucketState.BucketReferenced, BtnValidation := bench.Operator.JoyBtnRaw);
ADVANCE_TIME(10000000);
bench(M1_PresetTriggerCmd := encoderM1.HwOut.PresetTriggerCmd, M1_PresetValueOut := encoderM1.HwOut.PresetValueOut, M2_PresetTriggerCmd := encoderM2.HwOut.PresetTriggerCmd, M2_PresetValueOut := encoderM2.HwOut.PresetValueOut, RawPosM1 := raw1, RawPosM2 := raw2); raw1 := bench.RawPosM1; raw2 := bench.RawPosM2;
hw1.RawPosIn := bench.Winch.COD1_PosValue; hw1.SlaveOperational := TRUE; hw2.RawPosIn := bench.Winch.COD2_PosValue; hw2.SlaveOperational := TRUE;
encoderM1(Enable := TRUE, HomingPermit := TRUE, HomingAtTargetM := btnM1, CfgHomingTargetM := 8.7, CfgTopSensorPosM := 8.7, HwIn := hw1, Cfg := cfgEncoder, Calib := calibM1); calibM1 := encoderM1.Calib;
bucketEdge(CLK := btnBucket);
encoderM2(Enable := TRUE, HomingPermit := TRUE, HomingAtTargetM := btnM2 OR bucketEdge.Q, CfgHomingTargetM := 23.7, CfgTopSensorPosM := 23.7, UseDynamicTarget := bucketEdge.Q, DynamicHomingTargetM := encoderM1.Measurement.CablePosM + cfgBucket.OffsetCloseM, HwIn := hw2, Cfg := cfgEncoder, Calib := calibM2); calibM2 := encoderM2.Calib;
bucket(Enable := TRUE, Mode := E_Mode.MAINT_N2, PowerContactorEngaged := TRUE, CablePosM1 := encoderM1.Measurement.CablePosM, CablePosM2 := encoderM2.Measurement.CablePosM, HomedM1 := encoderM1.Homed, HomedM2 := encoderM2.Homed, HomedAndReliableM1 := encoderM1.HomedAndReliable, HomedAndReliableM2 := encoderM2.HomedAndReliable, HomingSuspectM1 := encoderM1.HomingSuspect, HomingSuspectM2 := encoderM2.HomingSuspect, ConfirmClosePosition := btnBucket, Config := cfgBucket, BucketState := bucketState); bucketState := bucket.BucketState;
home.M1Status.HomedAndReliable := encoderM1.HomedAndReliable; home.M2Status.HomedAndReliable := encoderM2.HomedAndReliable; home(BucketOffsetValid := bucketState.BucketReferenced, BtnValidation := bench.Operator.JoyBtnRaw);
ADVANCE_TIME(10000000);
bench(M1_PresetTriggerCmd := encoderM1.HwOut.PresetTriggerCmd, M1_PresetValueOut := encoderM1.HwOut.PresetValueOut, M2_PresetTriggerCmd := encoderM2.HwOut.PresetTriggerCmd, M2_PresetValueOut := encoderM2.HwOut.PresetValueOut, RawPosM1 := raw1, RawPosM2 := raw2); raw1 := bench.RawPosM1; raw2 := bench.RawPosM2;
hw1.RawPosIn := bench.Winch.COD1_PosValue; hw1.SlaveOperational := TRUE; hw2.RawPosIn := bench.Winch.COD2_PosValue; hw2.SlaveOperational := TRUE;
encoderM1(Enable := TRUE, HomingPermit := TRUE, HomingAtTargetM := btnM1, CfgHomingTargetM := 8.7, CfgTopSensorPosM := 8.7, HwIn := hw1, Cfg := cfgEncoder, Calib := calibM1); calibM1 := encoderM1.Calib;
bucketEdge(CLK := btnBucket);
encoderM2(Enable := TRUE, HomingPermit := TRUE, HomingAtTargetM := btnM2 OR bucketEdge.Q, CfgHomingTargetM := 23.7, CfgTopSensorPosM := 23.7, UseDynamicTarget := bucketEdge.Q, DynamicHomingTargetM := encoderM1.Measurement.CablePosM + cfgBucket.OffsetCloseM, HwIn := hw2, Cfg := cfgEncoder, Calib := calibM2); calibM2 := encoderM2.Calib;
bucket(Enable := TRUE, Mode := E_Mode.MAINT_N2, PowerContactorEngaged := TRUE, CablePosM1 := encoderM1.Measurement.CablePosM, CablePosM2 := encoderM2.Measurement.CablePosM, HomedM1 := encoderM1.Homed, HomedM2 := encoderM2.Homed, HomedAndReliableM1 := encoderM1.HomedAndReliable, HomedAndReliableM2 := encoderM2.HomedAndReliable, HomingSuspectM1 := encoderM1.HomingSuspect, HomingSuspectM2 := encoderM2.HomingSuspect, ConfirmClosePosition := btnBucket, Config := cfgBucket, BucketState := bucketState); bucketState := bucket.BucketState;
home.M1Status.HomedAndReliable := encoderM1.HomedAndReliable; home.M2Status.HomedAndReliable := encoderM2.HomedAndReliable; home(BucketOffsetValid := bucketState.BucketReferenced, BtnValidation := bench.Operator.JoyBtnRaw);
ADVANCE_TIME(10000000);
bench(M1_PresetTriggerCmd := encoderM1.HwOut.PresetTriggerCmd, M1_PresetValueOut := encoderM1.HwOut.PresetValueOut, M2_PresetTriggerCmd := encoderM2.HwOut.PresetTriggerCmd, M2_PresetValueOut := encoderM2.HwOut.PresetValueOut, RawPosM1 := raw1, RawPosM2 := raw2); raw1 := bench.RawPosM1; raw2 := bench.RawPosM2;
hw1.RawPosIn := bench.Winch.COD1_PosValue; hw1.SlaveOperational := TRUE; hw2.RawPosIn := bench.Winch.COD2_PosValue; hw2.SlaveOperational := TRUE;
encoderM1(Enable := TRUE, HomingPermit := TRUE, HomingAtTargetM := btnM1, CfgHomingTargetM := 8.7, CfgTopSensorPosM := 8.7, HwIn := hw1, Cfg := cfgEncoder, Calib := calibM1); calibM1 := encoderM1.Calib;
bucketEdge(CLK := btnBucket);
encoderM2(Enable := TRUE, HomingPermit := TRUE, HomingAtTargetM := btnM2 OR bucketEdge.Q, CfgHomingTargetM := 23.7, CfgTopSensorPosM := 23.7, UseDynamicTarget := bucketEdge.Q, DynamicHomingTargetM := encoderM1.Measurement.CablePosM + cfgBucket.OffsetCloseM, HwIn := hw2, Cfg := cfgEncoder, Calib := calibM2); calibM2 := encoderM2.Calib;
bucket(Enable := TRUE, Mode := E_Mode.MAINT_N2, PowerContactorEngaged := TRUE, CablePosM1 := encoderM1.Measurement.CablePosM, CablePosM2 := encoderM2.Measurement.CablePosM, HomedM1 := encoderM1.Homed, HomedM2 := encoderM2.Homed, HomedAndReliableM1 := encoderM1.HomedAndReliable, HomedAndReliableM2 := encoderM2.HomedAndReliable, HomingSuspectM1 := encoderM1.HomingSuspect, HomingSuspectM2 := encoderM2.HomingSuspect, ConfirmClosePosition := btnBucket, Config := cfgBucket, BucketState := bucketState); bucketState := bucket.BucketState;
home.M1Status.HomedAndReliable := encoderM1.HomedAndReliable; home.M2Status.HomedAndReliable := encoderM2.HomedAndReliable; home(BucketOffsetValid := bucketState.BucketReferenced, BtnValidation := bench.Operator.JoyBtnRaw);
ADVANCE_TIME(10000000);
bench(M1_PresetTriggerCmd := encoderM1.HwOut.PresetTriggerCmd, M1_PresetValueOut := encoderM1.HwOut.PresetValueOut, M2_PresetTriggerCmd := encoderM2.HwOut.PresetTriggerCmd, M2_PresetValueOut := encoderM2.HwOut.PresetValueOut, RawPosM1 := raw1, RawPosM2 := raw2); raw1 := bench.RawPosM1; raw2 := bench.RawPosM2;
hw1.RawPosIn := bench.Winch.COD1_PosValue; hw1.SlaveOperational := TRUE; hw2.RawPosIn := bench.Winch.COD2_PosValue; hw2.SlaveOperational := TRUE;
encoderM1(Enable := TRUE, HomingPermit := TRUE, HomingAtTargetM := btnM1, CfgHomingTargetM := 8.7, CfgTopSensorPosM := 8.7, HwIn := hw1, Cfg := cfgEncoder, Calib := calibM1); calibM1 := encoderM1.Calib;
bucketEdge(CLK := btnBucket);
encoderM2(Enable := TRUE, HomingPermit := TRUE, HomingAtTargetM := btnM2 OR bucketEdge.Q, CfgHomingTargetM := 23.7, CfgTopSensorPosM := 23.7, UseDynamicTarget := bucketEdge.Q, DynamicHomingTargetM := encoderM1.Measurement.CablePosM + cfgBucket.OffsetCloseM, HwIn := hw2, Cfg := cfgEncoder, Calib := calibM2); calibM2 := encoderM2.Calib;
bucket(Enable := TRUE, Mode := E_Mode.MAINT_N2, PowerContactorEngaged := TRUE, CablePosM1 := encoderM1.Measurement.CablePosM, CablePosM2 := encoderM2.Measurement.CablePosM, HomedM1 := encoderM1.Homed, HomedM2 := encoderM2.Homed, HomedAndReliableM1 := encoderM1.HomedAndReliable, HomedAndReliableM2 := encoderM2.HomedAndReliable, HomingSuspectM1 := encoderM1.HomingSuspect, HomingSuspectM2 := encoderM2.HomingSuspect, ConfirmClosePosition := btnBucket, Config := cfgBucket, BucketState := bucketState); bucketState := bucket.BucketState;
home.M1Status.HomedAndReliable := encoderM1.HomedAndReliable; home.M2Status.HomedAndReliable := encoderM2.HomedAndReliable; home(BucketOffsetValid := bucketState.BucketReferenced, BtnValidation := bench.Operator.JoyBtnRaw);
ADVANCE_TIME(10000000);
bench(M1_PresetTriggerCmd := encoderM1.HwOut.PresetTriggerCmd, M1_PresetValueOut := encoderM1.HwOut.PresetValueOut, M2_PresetTriggerCmd := encoderM2.HwOut.PresetTriggerCmd, M2_PresetValueOut := encoderM2.HwOut.PresetValueOut, RawPosM1 := raw1, RawPosM2 := raw2); raw1 := bench.RawPosM1; raw2 := bench.RawPosM2;
hw1.RawPosIn := bench.Winch.COD1_PosValue; hw1.SlaveOperational := TRUE; hw2.RawPosIn := bench.Winch.COD2_PosValue; hw2.SlaveOperational := TRUE;
encoderM1(Enable := TRUE, HomingPermit := TRUE, HomingAtTargetM := btnM1, CfgHomingTargetM := 8.7, CfgTopSensorPosM := 8.7, HwIn := hw1, Cfg := cfgEncoder, Calib := calibM1); calibM1 := encoderM1.Calib;
bucketEdge(CLK := btnBucket);
encoderM2(Enable := TRUE, HomingPermit := TRUE, HomingAtTargetM := btnM2 OR bucketEdge.Q, CfgHomingTargetM := 23.7, CfgTopSensorPosM := 23.7, UseDynamicTarget := bucketEdge.Q, DynamicHomingTargetM := encoderM1.Measurement.CablePosM + cfgBucket.OffsetCloseM, HwIn := hw2, Cfg := cfgEncoder, Calib := calibM2); calibM2 := encoderM2.Calib;
bucket(Enable := TRUE, Mode := E_Mode.MAINT_N2, PowerContactorEngaged := TRUE, CablePosM1 := encoderM1.Measurement.CablePosM, CablePosM2 := encoderM2.Measurement.CablePosM, HomedM1 := encoderM1.Homed, HomedM2 := encoderM2.Homed, HomedAndReliableM1 := encoderM1.HomedAndReliable, HomedAndReliableM2 := encoderM2.HomedAndReliable, HomingSuspectM1 := encoderM1.HomingSuspect, HomingSuspectM2 := encoderM2.HomingSuspect, ConfirmClosePosition := btnBucket, Config := cfgBucket, BucketState := bucketState); bucketState := bucket.BucketState;
home.M1Status.HomedAndReliable := encoderM1.HomedAndReliable; home.M2Status.HomedAndReliable := encoderM2.HomedAndReliable; home(BucketOffsetValid := bucketState.BucketReferenced, BtnValidation := bench.Operator.JoyBtnRaw);
ADVANCE_TIME(10000000);
bench(M1_PresetTriggerCmd := encoderM1.HwOut.PresetTriggerCmd, M1_PresetValueOut := encoderM1.HwOut.PresetValueOut, M2_PresetTriggerCmd := encoderM2.HwOut.PresetTriggerCmd, M2_PresetValueOut := encoderM2.HwOut.PresetValueOut, RawPosM1 := raw1, RawPosM2 := raw2); raw1 := bench.RawPosM1; raw2 := bench.RawPosM2;
hw1.RawPosIn := bench.Winch.COD1_PosValue; hw1.SlaveOperational := TRUE; hw2.RawPosIn := bench.Winch.COD2_PosValue; hw2.SlaveOperational := TRUE;
encoderM1(Enable := TRUE, HomingPermit := TRUE, HomingAtTargetM := btnM1, CfgHomingTargetM := 8.7, CfgTopSensorPosM := 8.7, HwIn := hw1, Cfg := cfgEncoder, Calib := calibM1); calibM1 := encoderM1.Calib;
bucketEdge(CLK := btnBucket);
encoderM2(Enable := TRUE, HomingPermit := TRUE, HomingAtTargetM := btnM2 OR bucketEdge.Q, CfgHomingTargetM := 23.7, CfgTopSensorPosM := 23.7, UseDynamicTarget := bucketEdge.Q, DynamicHomingTargetM := encoderM1.Measurement.CablePosM + cfgBucket.OffsetCloseM, HwIn := hw2, Cfg := cfgEncoder, Calib := calibM2); calibM2 := encoderM2.Calib;
bucket(Enable := TRUE, Mode := E_Mode.MAINT_N2, PowerContactorEngaged := TRUE, CablePosM1 := encoderM1.Measurement.CablePosM, CablePosM2 := encoderM2.Measurement.CablePosM, HomedM1 := encoderM1.Homed, HomedM2 := encoderM2.Homed, HomedAndReliableM1 := encoderM1.HomedAndReliable, HomedAndReliableM2 := encoderM2.HomedAndReliable, HomingSuspectM1 := encoderM1.HomingSuspect, HomingSuspectM2 := encoderM2.HomingSuspect, ConfirmClosePosition := btnBucket, Config := cfgBucket, BucketState := bucketState); bucketState := bucket.BucketState;
home.M1Status.HomedAndReliable := encoderM1.HomedAndReliable; home.M2Status.HomedAndReliable := encoderM2.HomedAndReliable; home(BucketOffsetValid := bucketState.BucketReferenced, BtnValidation := bench.Operator.JoyBtnRaw);
ADVANCE_TIME(10000000);
bench(M1_PresetTriggerCmd := encoderM1.HwOut.PresetTriggerCmd, M1_PresetValueOut := encoderM1.HwOut.PresetValueOut, M2_PresetTriggerCmd := encoderM2.HwOut.PresetTriggerCmd, M2_PresetValueOut := encoderM2.HwOut.PresetValueOut, RawPosM1 := raw1, RawPosM2 := raw2); raw1 := bench.RawPosM1; raw2 := bench.RawPosM2;
hw1.RawPosIn := bench.Winch.COD1_PosValue; hw1.SlaveOperational := TRUE; hw2.RawPosIn := bench.Winch.COD2_PosValue; hw2.SlaveOperational := TRUE;
encoderM1(Enable := TRUE, HomingPermit := TRUE, HomingAtTargetM := btnM1, CfgHomingTargetM := 8.7, CfgTopSensorPosM := 8.7, HwIn := hw1, Cfg := cfgEncoder, Calib := calibM1); calibM1 := encoderM1.Calib;
bucketEdge(CLK := btnBucket);
encoderM2(Enable := TRUE, HomingPermit := TRUE, HomingAtTargetM := btnM2 OR bucketEdge.Q, CfgHomingTargetM := 23.7, CfgTopSensorPosM := 23.7, UseDynamicTarget := bucketEdge.Q, DynamicHomingTargetM := encoderM1.Measurement.CablePosM + cfgBucket.OffsetCloseM, HwIn := hw2, Cfg := cfgEncoder, Calib := calibM2); calibM2 := encoderM2.Calib;
bucket(Enable := TRUE, Mode := E_Mode.MAINT_N2, PowerContactorEngaged := TRUE, CablePosM1 := encoderM1.Measurement.CablePosM, CablePosM2 := encoderM2.Measurement.CablePosM, HomedM1 := encoderM1.Homed, HomedM2 := encoderM2.Homed, HomedAndReliableM1 := encoderM1.HomedAndReliable, HomedAndReliableM2 := encoderM2.HomedAndReliable, HomingSuspectM1 := encoderM1.HomingSuspect, HomingSuspectM2 := encoderM2.HomingSuspect, ConfirmClosePosition := btnBucket, Config := cfgBucket, BucketState := bucketState); bucketState := bucket.BucketState;
home.M1Status.HomedAndReliable := encoderM1.HomedAndReliable; home.M2Status.HomedAndReliable := encoderM2.HomedAndReliable; home(BucketOffsetValid := bucketState.BucketReferenced, BtnValidation := bench.Operator.JoyBtnRaw);
ADVANCE_TIME(10000000);
bench(M1_PresetTriggerCmd := encoderM1.HwOut.PresetTriggerCmd, M1_PresetValueOut := encoderM1.HwOut.PresetValueOut, M2_PresetTriggerCmd := encoderM2.HwOut.PresetTriggerCmd, M2_PresetValueOut := encoderM2.HwOut.PresetValueOut, RawPosM1 := raw1, RawPosM2 := raw2); raw1 := bench.RawPosM1; raw2 := bench.RawPosM2;
hw1.RawPosIn := bench.Winch.COD1_PosValue; hw1.SlaveOperational := TRUE; hw2.RawPosIn := bench.Winch.COD2_PosValue; hw2.SlaveOperational := TRUE;
encoderM1(Enable := TRUE, HomingPermit := TRUE, HomingAtTargetM := btnM1, CfgHomingTargetM := 8.7, CfgTopSensorPosM := 8.7, HwIn := hw1, Cfg := cfgEncoder, Calib := calibM1); calibM1 := encoderM1.Calib;
bucketEdge(CLK := btnBucket);
encoderM2(Enable := TRUE, HomingPermit := TRUE, HomingAtTargetM := btnM2 OR bucketEdge.Q, CfgHomingTargetM := 23.7, CfgTopSensorPosM := 23.7, UseDynamicTarget := bucketEdge.Q, DynamicHomingTargetM := encoderM1.Measurement.CablePosM + cfgBucket.OffsetCloseM, HwIn := hw2, Cfg := cfgEncoder, Calib := calibM2); calibM2 := encoderM2.Calib;
bucket(Enable := TRUE, Mode := E_Mode.MAINT_N2, PowerContactorEngaged := TRUE, CablePosM1 := encoderM1.Measurement.CablePosM, CablePosM2 := encoderM2.Measurement.CablePosM, HomedM1 := encoderM1.Homed, HomedM2 := encoderM2.Homed, HomedAndReliableM1 := encoderM1.HomedAndReliable, HomedAndReliableM2 := encoderM2.HomedAndReliable, HomingSuspectM1 := encoderM1.HomingSuspect, HomingSuspectM2 := encoderM2.HomingSuspect, ConfirmClosePosition := btnBucket, Config := cfgBucket, BucketState := bucketState); bucketState := bucket.BucketState;
home.M1Status.HomedAndReliable := encoderM1.HomedAndReliable; home.M2Status.HomedAndReliable := encoderM2.HomedAndReliable; home(BucketOffsetValid := bucketState.BucketReferenced, BtnValidation := bench.Operator.JoyBtnRaw);
ADVANCE_TIME(10000000);
bench(M1_PresetTriggerCmd := encoderM1.HwOut.PresetTriggerCmd, M1_PresetValueOut := encoderM1.HwOut.PresetValueOut, M2_PresetTriggerCmd := encoderM2.HwOut.PresetTriggerCmd, M2_PresetValueOut := encoderM2.HwOut.PresetValueOut, RawPosM1 := raw1, RawPosM2 := raw2); raw1 := bench.RawPosM1; raw2 := bench.RawPosM2;
hw1.RawPosIn := bench.Winch.COD1_PosValue; hw1.SlaveOperational := TRUE; hw2.RawPosIn := bench.Winch.COD2_PosValue; hw2.SlaveOperational := TRUE;
encoderM1(Enable := TRUE, HomingPermit := TRUE, HomingAtTargetM := btnM1, CfgHomingTargetM := 8.7, CfgTopSensorPosM := 8.7, HwIn := hw1, Cfg := cfgEncoder, Calib := calibM1); calibM1 := encoderM1.Calib;
bucketEdge(CLK := btnBucket);
encoderM2(Enable := TRUE, HomingPermit := TRUE, HomingAtTargetM := btnM2 OR bucketEdge.Q, CfgHomingTargetM := 23.7, CfgTopSensorPosM := 23.7, UseDynamicTarget := bucketEdge.Q, DynamicHomingTargetM := encoderM1.Measurement.CablePosM + cfgBucket.OffsetCloseM, HwIn := hw2, Cfg := cfgEncoder, Calib := calibM2); calibM2 := encoderM2.Calib;
bucket(Enable := TRUE, Mode := E_Mode.MAINT_N2, PowerContactorEngaged := TRUE, CablePosM1 := encoderM1.Measurement.CablePosM, CablePosM2 := encoderM2.Measurement.CablePosM, HomedM1 := encoderM1.Homed, HomedM2 := encoderM2.Homed, HomedAndReliableM1 := encoderM1.HomedAndReliable, HomedAndReliableM2 := encoderM2.HomedAndReliable, HomingSuspectM1 := encoderM1.HomingSuspect, HomingSuspectM2 := encoderM2.HomingSuspect, ConfirmClosePosition := btnBucket, Config := cfgBucket, BucketState := bucketState); bucketState := bucket.BucketState;
home.M1Status.HomedAndReliable := encoderM1.HomedAndReliable; home.M2Status.HomedAndReliable := encoderM2.HomedAndReliable; home(BucketOffsetValid := bucketState.BucketReferenced, BtnValidation := bench.Operator.JoyBtnRaw);
ADVANCE_TIME(10000000);
bench(M1_PresetTriggerCmd := encoderM1.HwOut.PresetTriggerCmd, M1_PresetValueOut := encoderM1.HwOut.PresetValueOut, M2_PresetTriggerCmd := encoderM2.HwOut.PresetTriggerCmd, M2_PresetValueOut := encoderM2.HwOut.PresetValueOut, RawPosM1 := raw1, RawPosM2 := raw2); raw1 := bench.RawPosM1; raw2 := bench.RawPosM2;
hw1.RawPosIn := bench.Winch.COD1_PosValue; hw1.SlaveOperational := TRUE; hw2.RawPosIn := bench.Winch.COD2_PosValue; hw2.SlaveOperational := TRUE;
encoderM1(Enable := TRUE, HomingPermit := TRUE, HomingAtTargetM := btnM1, CfgHomingTargetM := 8.7, CfgTopSensorPosM := 8.7, HwIn := hw1, Cfg := cfgEncoder, Calib := calibM1); calibM1 := encoderM1.Calib;
bucketEdge(CLK := btnBucket);
encoderM2(Enable := TRUE, HomingPermit := TRUE, HomingAtTargetM := btnM2 OR bucketEdge.Q, CfgHomingTargetM := 23.7, CfgTopSensorPosM := 23.7, UseDynamicTarget := bucketEdge.Q, DynamicHomingTargetM := encoderM1.Measurement.CablePosM + cfgBucket.OffsetCloseM, HwIn := hw2, Cfg := cfgEncoder, Calib := calibM2); calibM2 := encoderM2.Calib;
bucket(Enable := TRUE, Mode := E_Mode.MAINT_N2, PowerContactorEngaged := TRUE, CablePosM1 := encoderM1.Measurement.CablePosM, CablePosM2 := encoderM2.Measurement.CablePosM, HomedM1 := encoderM1.Homed, HomedM2 := encoderM2.Homed, HomedAndReliableM1 := encoderM1.HomedAndReliable, HomedAndReliableM2 := encoderM2.HomedAndReliable, HomingSuspectM1 := encoderM1.HomingSuspect, HomingSuspectM2 := encoderM2.HomingSuspect, ConfirmClosePosition := btnBucket, Config := cfgBucket, BucketState := bucketState); bucketState := bucket.BucketState;
home.M1Status.HomedAndReliable := encoderM1.HomedAndReliable; home.M2Status.HomedAndReliable := encoderM2.HomedAndReliable; home(BucketOffsetValid := bucketState.BucketReferenced, BtnValidation := bench.Operator.JoyBtnRaw);
ADVANCE_TIME(10000000);
bench(M1_PresetTriggerCmd := encoderM1.HwOut.PresetTriggerCmd, M1_PresetValueOut := encoderM1.HwOut.PresetValueOut, M2_PresetTriggerCmd := encoderM2.HwOut.PresetTriggerCmd, M2_PresetValueOut := encoderM2.HwOut.PresetValueOut, RawPosM1 := raw1, RawPosM2 := raw2); raw1 := bench.RawPosM1; raw2 := bench.RawPosM2;
hw1.RawPosIn := bench.Winch.COD1_PosValue; hw1.SlaveOperational := TRUE; hw2.RawPosIn := bench.Winch.COD2_PosValue; hw2.SlaveOperational := TRUE;
encoderM1(Enable := TRUE, HomingPermit := TRUE, HomingAtTargetM := btnM1, CfgHomingTargetM := 8.7, CfgTopSensorPosM := 8.7, HwIn := hw1, Cfg := cfgEncoder, Calib := calibM1); calibM1 := encoderM1.Calib;
bucketEdge(CLK := btnBucket);
encoderM2(Enable := TRUE, HomingPermit := TRUE, HomingAtTargetM := btnM2 OR bucketEdge.Q, CfgHomingTargetM := 23.7, CfgTopSensorPosM := 23.7, UseDynamicTarget := bucketEdge.Q, DynamicHomingTargetM := encoderM1.Measurement.CablePosM + cfgBucket.OffsetCloseM, HwIn := hw2, Cfg := cfgEncoder, Calib := calibM2); calibM2 := encoderM2.Calib;
bucket(Enable := TRUE, Mode := E_Mode.MAINT_N2, PowerContactorEngaged := TRUE, CablePosM1 := encoderM1.Measurement.CablePosM, CablePosM2 := encoderM2.Measurement.CablePosM, HomedM1 := encoderM1.Homed, HomedM2 := encoderM2.Homed, HomedAndReliableM1 := encoderM1.HomedAndReliable, HomedAndReliableM2 := encoderM2.HomedAndReliable, HomingSuspectM1 := encoderM1.HomingSuspect, HomingSuspectM2 := encoderM2.HomingSuspect, ConfirmClosePosition := btnBucket, Config := cfgBucket, BucketState := bucketState); bucketState := bucket.BucketState;
home.M1Status.HomedAndReliable := encoderM1.HomedAndReliable; home.M2Status.HomedAndReliable := encoderM2.HomedAndReliable; home(BucketOffsetValid := bucketState.BucketReferenced, BtnValidation := bench.Operator.JoyBtnRaw);
ADVANCE_TIME(10000000);
bench(M1_PresetTriggerCmd := encoderM1.HwOut.PresetTriggerCmd, M1_PresetValueOut := encoderM1.HwOut.PresetValueOut, M2_PresetTriggerCmd := encoderM2.HwOut.PresetTriggerCmd, M2_PresetValueOut := encoderM2.HwOut.PresetValueOut, RawPosM1 := raw1, RawPosM2 := raw2); raw1 := bench.RawPosM1; raw2 := bench.RawPosM2;
hw1.RawPosIn := bench.Winch.COD1_PosValue; hw1.SlaveOperational := TRUE; hw2.RawPosIn := bench.Winch.COD2_PosValue; hw2.SlaveOperational := TRUE;
encoderM1(Enable := TRUE, HomingPermit := TRUE, HomingAtTargetM := btnM1, CfgHomingTargetM := 8.7, CfgTopSensorPosM := 8.7, HwIn := hw1, Cfg := cfgEncoder, Calib := calibM1); calibM1 := encoderM1.Calib;
bucketEdge(CLK := btnBucket);
encoderM2(Enable := TRUE, HomingPermit := TRUE, HomingAtTargetM := btnM2 OR bucketEdge.Q, CfgHomingTargetM := 23.7, CfgTopSensorPosM := 23.7, UseDynamicTarget := bucketEdge.Q, DynamicHomingTargetM := encoderM1.Measurement.CablePosM + cfgBucket.OffsetCloseM, HwIn := hw2, Cfg := cfgEncoder, Calib := calibM2); calibM2 := encoderM2.Calib;
bucket(Enable := TRUE, Mode := E_Mode.MAINT_N2, PowerContactorEngaged := TRUE, CablePosM1 := encoderM1.Measurement.CablePosM, CablePosM2 := encoderM2.Measurement.CablePosM, HomedM1 := encoderM1.Homed, HomedM2 := encoderM2.Homed, HomedAndReliableM1 := encoderM1.HomedAndReliable, HomedAndReliableM2 := encoderM2.HomedAndReliable, HomingSuspectM1 := encoderM1.HomingSuspect, HomingSuspectM2 := encoderM2.HomingSuspect, ConfirmClosePosition := btnBucket, Config := cfgBucket, BucketState := bucketState); bucketState := bucket.BucketState;
home.M1Status.HomedAndReliable := encoderM1.HomedAndReliable; home.M2Status.HomedAndReliable := encoderM2.HomedAndReliable; home(BucketOffsetValid := bucketState.BucketReferenced, BtnValidation := bench.Operator.JoyBtnRaw);
ADVANCE_TIME(10000000);
bench(M1_PresetTriggerCmd := encoderM1.HwOut.PresetTriggerCmd, M1_PresetValueOut := encoderM1.HwOut.PresetValueOut, M2_PresetTriggerCmd := encoderM2.HwOut.PresetTriggerCmd, M2_PresetValueOut := encoderM2.HwOut.PresetValueOut, RawPosM1 := raw1, RawPosM2 := raw2); raw1 := bench.RawPosM1; raw2 := bench.RawPosM2;
hw1.RawPosIn := bench.Winch.COD1_PosValue; hw1.SlaveOperational := TRUE; hw2.RawPosIn := bench.Winch.COD2_PosValue; hw2.SlaveOperational := TRUE;
encoderM1(Enable := TRUE, HomingPermit := TRUE, HomingAtTargetM := btnM1, CfgHomingTargetM := 8.7, CfgTopSensorPosM := 8.7, HwIn := hw1, Cfg := cfgEncoder, Calib := calibM1); calibM1 := encoderM1.Calib;
bucketEdge(CLK := btnBucket);
encoderM2(Enable := TRUE, HomingPermit := TRUE, HomingAtTargetM := btnM2 OR bucketEdge.Q, CfgHomingTargetM := 23.7, CfgTopSensorPosM := 23.7, UseDynamicTarget := bucketEdge.Q, DynamicHomingTargetM := encoderM1.Measurement.CablePosM + cfgBucket.OffsetCloseM, HwIn := hw2, Cfg := cfgEncoder, Calib := calibM2); calibM2 := encoderM2.Calib;
bucket(Enable := TRUE, Mode := E_Mode.MAINT_N2, PowerContactorEngaged := TRUE, CablePosM1 := encoderM1.Measurement.CablePosM, CablePosM2 := encoderM2.Measurement.CablePosM, HomedM1 := encoderM1.Homed, HomedM2 := encoderM2.Homed, HomedAndReliableM1 := encoderM1.HomedAndReliable, HomedAndReliableM2 := encoderM2.HomedAndReliable, HomingSuspectM1 := encoderM1.HomingSuspect, HomingSuspectM2 := encoderM2.HomingSuspect, ConfirmClosePosition := btnBucket, Config := cfgBucket, BucketState := bucketState); bucketState := bucket.BucketState;
home.M1Status.HomedAndReliable := encoderM1.HomedAndReliable; home.M2Status.HomedAndReliable := encoderM2.HomedAndReliable; home(BucketOffsetValid := bucketState.BucketReferenced, BtnValidation := bench.Operator.JoyBtnRaw);
ADVANCE_TIME(10000000);
bench(M1_PresetTriggerCmd := encoderM1.HwOut.PresetTriggerCmd, M1_PresetValueOut := encoderM1.HwOut.PresetValueOut, M2_PresetTriggerCmd := encoderM2.HwOut.PresetTriggerCmd, M2_PresetValueOut := encoderM2.HwOut.PresetValueOut, RawPosM1 := raw1, RawPosM2 := raw2); raw1 := bench.RawPosM1; raw2 := bench.RawPosM2;
hw1.RawPosIn := bench.Winch.COD1_PosValue; hw1.SlaveOperational := TRUE; hw2.RawPosIn := bench.Winch.COD2_PosValue; hw2.SlaveOperational := TRUE;
encoderM1(Enable := TRUE, HomingPermit := TRUE, HomingAtTargetM := btnM1, CfgHomingTargetM := 8.7, CfgTopSensorPosM := 8.7, HwIn := hw1, Cfg := cfgEncoder, Calib := calibM1); calibM1 := encoderM1.Calib;
bucketEdge(CLK := btnBucket);
encoderM2(Enable := TRUE, HomingPermit := TRUE, HomingAtTargetM := btnM2 OR bucketEdge.Q, CfgHomingTargetM := 23.7, CfgTopSensorPosM := 23.7, UseDynamicTarget := bucketEdge.Q, DynamicHomingTargetM := encoderM1.Measurement.CablePosM + cfgBucket.OffsetCloseM, HwIn := hw2, Cfg := cfgEncoder, Calib := calibM2); calibM2 := encoderM2.Calib;
bucket(Enable := TRUE, Mode := E_Mode.MAINT_N2, PowerContactorEngaged := TRUE, CablePosM1 := encoderM1.Measurement.CablePosM, CablePosM2 := encoderM2.Measurement.CablePosM, HomedM1 := encoderM1.Homed, HomedM2 := encoderM2.Homed, HomedAndReliableM1 := encoderM1.HomedAndReliable, HomedAndReliableM2 := encoderM2.HomedAndReliable, HomingSuspectM1 := encoderM1.HomingSuspect, HomingSuspectM2 := encoderM2.HomingSuspect, ConfirmClosePosition := btnBucket, Config := cfgBucket, BucketState := bucketState); bucketState := bucket.BucketState;
home.M1Status.HomedAndReliable := encoderM1.HomedAndReliable; home.M2Status.HomedAndReliable := encoderM2.HomedAndReliable; home(BucketOffsetValid := bucketState.BucketReferenced, BtnValidation := bench.Operator.JoyBtnRaw);
ASSERT_TRUE(bucketState.BucketReferenced, 'Troisieme bouton confirme datum benne'); ASSERT_TRUE(home.MachineHomed, 'Qualification machine issue des vrais composants'); ASSERT_EQ(home.MachineHomingSeqStep, E_MachineHomingTxState.HX0_REPOS, 'Aucun lancement grafcet par references manuelles'); ASSERT_FALSE(home.M3Locked, 'Aucun verrou homing parasite');
END_TEST
